(* IEC 61131-3 sources: STAR-PLC-Agent/results/raw/codex_matrix_resume_20261114/codex_deepseek/PUB019/functional/attempt_0001, 1 file *)

(* ---- test_program.st ---- *)
PROGRAM PLC_PRG
VAR
 BenchStep : UDINT := 0;
 BenchCalls : UDINT := 0;
 BenchDone : BOOL := FALSE;
 BenchUut0 : FB_Task;
 BenchUut1 : FB_Task;
 BenchUut2 : FB_Task;
 BenchUut3 : FB_Task;
 BenchUut4 : FB_Task;
 BenchUut5 : FB_Task;
 BenchUut6 : FB_Task;
 BenchUut7 : FB_Task;
 BenchUut8 : FB_Task;
 BenchUut9 : FB_Task;
 BenchUut10 : FB_Task;
 BenchUut11 : FB_Task;
 BenchUut12 : FB_Task;
 BenchUut13 : FB_Task;
 BenchUut14 : FB_Task;
 BenchUut15 : FB_Task;
 BenchUut16 : FB_Task;
 TraceIn_ManualMode : ARRAY[0..305] OF BOOL;
 TraceIn_SingleStepMode : ARRAY[0..305] OF BOOL;
 TraceIn_SingleCycleMode : ARRAY[0..305] OF BOOL;
 TraceIn_ContinuousMode : ARRAY[0..305] OF BOOL;
 TraceIn_EmergencyStop : ARRAY[0..305] OF BOOL;
 TraceIn_Start : ARRAY[0..305] OF BOOL;
 TraceIn_DownButton : ARRAY[0..305] OF BOOL;
 TraceIn_UpButton : ARRAY[0..305] OF BOOL;
 TraceIn_LeftButton : ARRAY[0..305] OF BOOL;
 TraceIn_RightButton : ARRAY[0..305] OF BOOL;
 TraceIn_GripButton : ARRAY[0..305] OF BOOL;
 TraceIn_ReleaseButton : ARRAY[0..305] OF BOOL;
 TraceIn_DownLimitSwitch : ARRAY[0..305] OF BOOL;
 TraceIn_UpLimitSwitch : ARRAY[0..305] OF BOOL;
 TraceIn_LeftLimitSwitch : ARRAY[0..305] OF BOOL;
 TraceIn_RightLimitSwitch : ARRAY[0..305] OF BOOL;
 TraceIn_GripLimitSwitch : ARRAY[0..305] OF BOOL;
 TraceIn_ReleaseLimitSwitch : ARRAY[0..305] OF BOOL;
 TraceOut_MoveDown : ARRAY[0..305] OF BOOL;
 TraceOut_MoveUp : ARRAY[0..305] OF BOOL;
 TraceOut_MoveLeft : ARRAY[0..305] OF BOOL;
 TraceOut_MoveRight : ARRAY[0..305] OF BOOL;
 TraceOut_ActivateGrip : ARRAY[0..305] OF BOOL;
 TraceOut_ActivateRelease : ARRAY[0..305] OF BOOL;
END_VAR

IF NOT BenchDone THEN
 CASE BenchStep OF
 0:
   BenchUut0.ManualMode := TRUE;
   BenchUut0.SingleStepMode := FALSE;
   BenchUut0.SingleCycleMode := FALSE;
   BenchUut0.ContinuousMode := FALSE;
   BenchUut0.EmergencyStop := TRUE;
   BenchUut0.Start := FALSE;
   BenchUut0.DownButton := TRUE;
   BenchUut0.UpButton := FALSE;
   BenchUut0.LeftButton := FALSE;
   BenchUut0.RightButton := FALSE;
   BenchUut0.GripButton := FALSE;
   BenchUut0.ReleaseButton := FALSE;
   BenchUut0.DownLimitSwitch := FALSE;
   BenchUut0.UpLimitSwitch := TRUE;
   BenchUut0.LeftLimitSwitch := TRUE;
   BenchUut0.RightLimitSwitch := FALSE;
   BenchUut0.GripLimitSwitch := FALSE;
   BenchUut0.ReleaseLimitSwitch := TRUE;
   TraceIn_ManualMode[0] := BenchUut0.ManualMode;
   TraceIn_SingleStepMode[0] := BenchUut0.SingleStepMode;
   TraceIn_SingleCycleMode[0] := BenchUut0.SingleCycleMode;
   TraceIn_ContinuousMode[0] := BenchUut0.ContinuousMode;
   TraceIn_EmergencyStop[0] := BenchUut0.EmergencyStop;
   TraceIn_Start[0] := BenchUut0.Start;
   TraceIn_DownButton[0] := BenchUut0.DownButton;
   TraceIn_UpButton[0] := BenchUut0.UpButton;
   TraceIn_LeftButton[0] := BenchUut0.LeftButton;
   TraceIn_RightButton[0] := BenchUut0.RightButton;
   TraceIn_GripButton[0] := BenchUut0.GripButton;
   TraceIn_ReleaseButton[0] := BenchUut0.ReleaseButton;
   TraceIn_DownLimitSwitch[0] := BenchUut0.DownLimitSwitch;
   TraceIn_UpLimitSwitch[0] := BenchUut0.UpLimitSwitch;
   TraceIn_LeftLimitSwitch[0] := BenchUut0.LeftLimitSwitch;
   TraceIn_RightLimitSwitch[0] := BenchUut0.RightLimitSwitch;
   TraceIn_GripLimitSwitch[0] := BenchUut0.GripLimitSwitch;
   TraceIn_ReleaseLimitSwitch[0] := BenchUut0.ReleaseLimitSwitch;
   BenchUut0();
   TraceOut_MoveDown[0] := BenchUut0.MoveDown;
   TraceOut_MoveUp[0] := BenchUut0.MoveUp;
   TraceOut_MoveLeft[0] := BenchUut0.MoveLeft;
   TraceOut_MoveRight[0] := BenchUut0.MoveRight;
   TraceOut_ActivateGrip[0] := BenchUut0.ActivateGrip;
   TraceOut_ActivateRelease[0] := BenchUut0.ActivateRelease;
   BenchCalls := BenchCalls + 1;
 1:
   BenchUut0.ManualMode := TRUE;
   BenchUut0.SingleStepMode := FALSE;
   BenchUut0.SingleCycleMode := FALSE;
   BenchUut0.ContinuousMode := FALSE;
   BenchUut0.EmergencyStop := TRUE;
   BenchUut0.Start := FALSE;
   BenchUut0.DownButton := TRUE;
   BenchUut0.UpButton := FALSE;
   BenchUut0.LeftButton := FALSE;
   BenchUut0.RightButton := FALSE;
   BenchUut0.GripButton := FALSE;
   BenchUut0.ReleaseButton := FALSE;
   BenchUut0.DownLimitSwitch := TRUE;
   BenchUut0.UpLimitSwitch := FALSE;
   BenchUut0.LeftLimitSwitch := TRUE;
   BenchUut0.RightLimitSwitch := FALSE;
   BenchUut0.GripLimitSwitch := FALSE;
   BenchUut0.ReleaseLimitSwitch := TRUE;
   TraceIn_ManualMode[1] := BenchUut0.ManualMode;
   TraceIn_SingleStepMode[1] := BenchUut0.SingleStepMode;
   TraceIn_SingleCycleMode[1] := BenchUut0.SingleCycleMode;
   TraceIn_ContinuousMode[1] := BenchUut0.ContinuousMode;
   TraceIn_EmergencyStop[1] := BenchUut0.EmergencyStop;
   TraceIn_Start[1] := BenchUut0.Start;
   TraceIn_DownButton[1] := BenchUut0.DownButton;
   TraceIn_UpButton[1] := BenchUut0.UpButton;
   TraceIn_LeftButton[1] := BenchUut0.LeftButton;
   TraceIn_RightButton[1] := BenchUut0.RightButton;
   TraceIn_GripButton[1] := BenchUut0.GripButton;
   TraceIn_ReleaseButton[1] := BenchUut0.ReleaseButton;
   TraceIn_DownLimitSwitch[1] := BenchUut0.DownLimitSwitch;
   TraceIn_UpLimitSwitch[1] := BenchUut0.UpLimitSwitch;
   TraceIn_LeftLimitSwitch[1] := BenchUut0.LeftLimitSwitch;
   TraceIn_RightLimitSwitch[1] := BenchUut0.RightLimitSwitch;
   TraceIn_GripLimitSwitch[1] := BenchUut0.GripLimitSwitch;
   TraceIn_ReleaseLimitSwitch[1] := BenchUut0.ReleaseLimitSwitch;
   BenchUut0();
   TraceOut_MoveDown[1] := BenchUut0.MoveDown;
   TraceOut_MoveUp[1] := BenchUut0.MoveUp;
   TraceOut_MoveLeft[1] := BenchUut0.MoveLeft;
   TraceOut_MoveRight[1] := BenchUut0.MoveRight;
   TraceOut_ActivateGrip[1] := BenchUut0.ActivateGrip;
   TraceOut_ActivateRelease[1] := BenchUut0.ActivateRelease;
   BenchCalls := BenchCalls + 1;
 2:
   BenchUut0.ManualMode := TRUE;
   BenchUut0.SingleStepMode := FALSE;
   BenchUut0.SingleCycleMode := FALSE;
   BenchUut0.ContinuousMode := FALSE;
   BenchUut0.EmergencyStop := TRUE;
   BenchUut0.Start := FALSE;
   BenchUut0.DownButton := FALSE;
   BenchUut0.UpButton := FALSE;
   BenchUut0.LeftButton := FALSE;
   BenchUut0.RightButton := FALSE;
   BenchUut0.GripButton := FALSE;
   BenchUut0.ReleaseButton := FALSE;
   BenchUut0.DownLimitSwitch := FALSE;
   BenchUut0.UpLimitSwitch := TRUE;
   BenchUut0.LeftLimitSwitch := TRUE;
   BenchUut0.RightLimitSwitch := FALSE;
   BenchUut0.GripLimitSwitch := FALSE;
   BenchUut0.ReleaseLimitSwitch := TRUE;
   TraceIn_ManualMode[2] := BenchUut0.ManualMode;
   TraceIn_SingleStepMode[2] := BenchUut0.SingleStepMode;
   TraceIn_SingleCycleMode[2] := BenchUut0.SingleCycleMode;
   TraceIn_ContinuousMode[2] := BenchUut0.ContinuousMode;
   TraceIn_EmergencyStop[2] := BenchUut0.EmergencyStop;
   TraceIn_Start[2] := BenchUut0.Start;
   TraceIn_DownButton[2] := BenchUut0.DownButton;
   TraceIn_UpButton[2] := BenchUut0.UpButton;
   TraceIn_LeftButton[2] := BenchUut0.LeftButton;
   TraceIn_RightButton[2] := BenchUut0.RightButton;
   TraceIn_GripButton[2] := BenchUut0.GripButton;
   TraceIn_ReleaseButton[2] := BenchUut0.ReleaseButton;
   TraceIn_DownLimitSwitch[2] := BenchUut0.DownLimitSwitch;
   TraceIn_UpLimitSwitch[2] := BenchUut0.UpLimitSwitch;
   TraceIn_LeftLimitSwitch[2] := BenchUut0.LeftLimitSwitch;
   TraceIn_RightLimitSwitch[2] := BenchUut0.RightLimitSwitch;
   TraceIn_GripLimitSwitch[2] := BenchUut0.GripLimitSwitch;
   TraceIn_ReleaseLimitSwitch[2] := BenchUut0.ReleaseLimitSwitch;
   BenchUut0();
   TraceOut_MoveDown[2] := BenchUut0.MoveDown;
   TraceOut_MoveUp[2] := BenchUut0.MoveUp;
   TraceOut_MoveLeft[2] := BenchUut0.MoveLeft;
   TraceOut_MoveRight[2] := BenchUut0.MoveRight;
   TraceOut_ActivateGrip[2] := BenchUut0.ActivateGrip;
   TraceOut_ActivateRelease[2] := BenchUut0.ActivateRelease;
   BenchCalls := BenchCalls + 1;
 3:
   BenchUut0.ManualMode := TRUE;
   BenchUut0.SingleStepMode := FALSE;
   BenchUut0.SingleCycleMode := FALSE;
   BenchUut0.ContinuousMode := FALSE;
   BenchUut0.EmergencyStop := TRUE;
   BenchUut0.Start := FALSE;
   BenchUut0.DownButton := TRUE;
   BenchUut0.UpButton := TRUE;
   BenchUut0.LeftButton := FALSE;
   BenchUut0.RightButton := FALSE;
   BenchUut0.GripButton := FALSE;
   BenchUut0.ReleaseButton := FALSE;
   BenchUut0.DownLimitSwitch := FALSE;
   BenchUut0.UpLimitSwitch := FALSE;
   BenchUut0.LeftLimitSwitch := TRUE;
   BenchUut0.RightLimitSwitch := FALSE;
   BenchUut0.GripLimitSwitch := FALSE;
   BenchUut0.ReleaseLimitSwitch := TRUE;
   TraceIn_ManualMode[3] := BenchUut0.ManualMode;
   TraceIn_SingleStepMode[3] := BenchUut0.SingleStepMode;
   TraceIn_SingleCycleMode[3] := BenchUut0.SingleCycleMode;
   TraceIn_ContinuousMode[3] := BenchUut0.ContinuousMode;
   TraceIn_EmergencyStop[3] := BenchUut0.EmergencyStop;
   TraceIn_Start[3] := BenchUut0.Start;
   TraceIn_DownButton[3] := BenchUut0.DownButton;
   TraceIn_UpButton[3] := BenchUut0.UpButton;
   TraceIn_LeftButton[3] := BenchUut0.LeftButton;
   TraceIn_RightButton[3] := BenchUut0.RightButton;
   TraceIn_GripButton[3] := BenchUut0.GripButton;
   TraceIn_ReleaseButton[3] := BenchUut0.ReleaseButton;
   TraceIn_DownLimitSwitch[3] := BenchUut0.DownLimitSwitch;
   TraceIn_UpLimitSwitch[3] := BenchUut0.UpLimitSwitch;
   TraceIn_LeftLimitSwitch[3] := BenchUut0.LeftLimitSwitch;
   TraceIn_RightLimitSwitch[3] := BenchUut0.RightLimitSwitch;
   TraceIn_GripLimitSwitch[3] := BenchUut0.GripLimitSwitch;
   TraceIn_ReleaseLimitSwitch[3] := BenchUut0.ReleaseLimitSwitch;
   BenchUut0();
   TraceOut_MoveDown[3] := BenchUut0.MoveDown;
   TraceOut_MoveUp[3] := BenchUut0.MoveUp;
   TraceOut_MoveLeft[3] := BenchUut0.MoveLeft;
   TraceOut_MoveRight[3] := BenchUut0.MoveRight;
   TraceOut_ActivateGrip[3] := BenchUut0.ActivateGrip;
   TraceOut_ActivateRelease[3] := BenchUut0.ActivateRelease;
   BenchCalls := BenchCalls + 1;
 4:
   BenchUut0.ManualMode := TRUE;
   BenchUut0.SingleStepMode := FALSE;
   BenchUut0.SingleCycleMode := FALSE;
   BenchUut0.ContinuousMode := FALSE;
   BenchUut0.EmergencyStop := TRUE;
   BenchUut0.Start := FALSE;
   BenchUut0.DownButton := FALSE;
   BenchUut0.UpButton := FALSE;
   BenchUut0.LeftButton := FALSE;
   BenchUut0.RightButton := TRUE;
   BenchUut0.GripButton := FALSE;
   BenchUut0.ReleaseButton := FALSE;
   BenchUut0.DownLimitSwitch := FALSE;
   BenchUut0.UpLimitSwitch := TRUE;
   BenchUut0.LeftLimitSwitch := TRUE;
   BenchUut0.RightLimitSwitch := FALSE;
   BenchUut0.GripLimitSwitch := FALSE;
   BenchUut0.ReleaseLimitSwitch := TRUE;
   TraceIn_ManualMode[4] := BenchUut0.ManualMode;
   TraceIn_SingleStepMode[4] := BenchUut0.SingleStepMode;
   TraceIn_SingleCycleMode[4] := BenchUut0.SingleCycleMode;
   TraceIn_ContinuousMode[4] := BenchUut0.ContinuousMode;
   TraceIn_EmergencyStop[4] := BenchUut0.EmergencyStop;
   TraceIn_Start[4] := BenchUut0.Start;
   TraceIn_DownButton[4] := BenchUut0.DownButton;
   TraceIn_UpButton[4] := BenchUut0.UpButton;
   TraceIn_LeftButton[4] := BenchUut0.LeftButton;
   TraceIn_RightButton[4] := BenchUut0.RightButton;
   TraceIn_GripButton[4] := BenchUut0.GripButton;
   TraceIn_ReleaseButton[4] := BenchUut0.ReleaseButton;
   TraceIn_DownLimitSwitch[4] := BenchUut0.DownLimitSwitch;
   TraceIn_UpLimitSwitch[4] := BenchUut0.UpLimitSwitch;
   TraceIn_LeftLimitSwitch[4] := BenchUut0.LeftLimitSwitch;
   TraceIn_RightLimitSwitch[4] := BenchUut0.RightLimitSwitch;
   TraceIn_GripLimitSwitch[4] := BenchUut0.GripLimitSwitch;
   TraceIn_ReleaseLimitSwitch[4] := BenchUut0.ReleaseLimitSwitch;
   BenchUut0();
   TraceOut_MoveDown[4] := BenchUut0.MoveDown;
   TraceOut_MoveUp[4] := BenchUut0.MoveUp;
   TraceOut_MoveLeft[4] := BenchUut0.MoveLeft;
   TraceOut_MoveRight[4] := BenchUut0.MoveRight;
   TraceOut_ActivateGrip[4] := BenchUut0.ActivateGrip;
   TraceOut_ActivateRelease[4] := BenchUut0.ActivateRelease;
   BenchCalls := BenchCalls + 1;
 5:
   BenchUut0.ManualMode := TRUE;
   BenchUut0.SingleStepMode := FALSE;
   BenchUut0.SingleCycleMode := FALSE;
   BenchUut0.ContinuousMode := FALSE;
   BenchUut0.EmergencyStop := TRUE;
   BenchUut0.Start := FALSE;
   BenchUut0.DownButton := FALSE;
   BenchUut0.UpButton := FALSE;
   BenchUut0.LeftButton := FALSE;
   BenchUut0.RightButton := TRUE;
   BenchUut0.GripButton := FALSE;
   BenchUut0.ReleaseButton := FALSE;
   BenchUut0.DownLimitSwitch := FALSE;
   BenchUut0.UpLimitSwitch := TRUE;
   BenchUut0.LeftLimitSwitch := FALSE;
   BenchUut0.RightLimitSwitch := TRUE;
   BenchUut0.GripLimitSwitch := FALSE;
   BenchUut0.ReleaseLimitSwitch := TRUE;
   TraceIn_ManualMode[5] := BenchUut0.ManualMode;
   TraceIn_SingleStepMode[5] := BenchUut0.SingleStepMode;
   TraceIn_SingleCycleMode[5] := BenchUut0.SingleCycleMode;
   TraceIn_ContinuousMode[5] := BenchUut0.ContinuousMode;
   TraceIn_EmergencyStop[5] := BenchUut0.EmergencyStop;
   TraceIn_Start[5] := BenchUut0.Start;
   TraceIn_DownButton[5] := BenchUut0.DownButton;
   TraceIn_UpButton[5] := BenchUut0.UpButton;
   TraceIn_LeftButton[5] := BenchUut0.LeftButton;
   TraceIn_RightButton[5] := BenchUut0.RightButton;
   TraceIn_GripButton[5] := BenchUut0.GripButton;
   TraceIn_ReleaseButton[5] := BenchUut0.ReleaseButton;
   TraceIn_DownLimitSwitch[5] := BenchUut0.DownLimitSwitch;
   TraceIn_UpLimitSwitch[5] := BenchUut0.UpLimitSwitch;
   TraceIn_LeftLimitSwitch[5] := BenchUut0.LeftLimitSwitch;
   TraceIn_RightLimitSwitch[5] := BenchUut0.RightLimitSwitch;
   TraceIn_GripLimitSwitch[5] := BenchUut0.GripLimitSwitch;
   TraceIn_ReleaseLimitSwitch[5] := BenchUut0.ReleaseLimitSwitch;
   BenchUut0();
   TraceOut_MoveDown[5] := BenchUut0.MoveDown;
   TraceOut_MoveUp[5] := BenchUut0.MoveUp;
   TraceOut_MoveLeft[5] := BenchUut0.MoveLeft;
   TraceOut_MoveRight[5] := BenchUut0.MoveRight;
   TraceOut_ActivateGrip[5] := BenchUut0.ActivateGrip;
   TraceOut_ActivateRelease[5] := BenchUut0.ActivateRelease;
   BenchCalls := BenchCalls + 1;
 6:
   BenchUut0.ManualMode := TRUE;
   BenchUut0.SingleStepMode := FALSE;
   BenchUut0.SingleCycleMode := FALSE;
   BenchUut0.ContinuousMode := FALSE;
   BenchUut0.EmergencyStop := TRUE;
   BenchUut0.Start := FALSE;
   BenchUut0.DownButton := FALSE;
   BenchUut0.UpButton := FALSE;
   BenchUut0.LeftButton := FALSE;
   BenchUut0.RightButton := FALSE;
   BenchUut0.GripButton := TRUE;
   BenchUut0.ReleaseButton := FALSE;
   BenchUut0.DownLimitSwitch := FALSE;
   BenchUut0.UpLimitSwitch := TRUE;
   BenchUut0.LeftLimitSwitch := TRUE;
   BenchUut0.RightLimitSwitch := FALSE;
   BenchUut0.GripLimitSwitch := FALSE;
   BenchUut0.ReleaseLimitSwitch := FALSE;
   TraceIn_ManualMode[6] := BenchUut0.ManualMode;
   TraceIn_SingleStepMode[6] := BenchUut0.SingleStepMode;
   TraceIn_SingleCycleMode[6] := BenchUut0.SingleCycleMode;
   TraceIn_ContinuousMode[6] := BenchUut0.ContinuousMode;
   TraceIn_EmergencyStop[6] := BenchUut0.EmergencyStop;
   TraceIn_Start[6] := BenchUut0.Start;
   TraceIn_DownButton[6] := BenchUut0.DownButton;
   TraceIn_UpButton[6] := BenchUut0.UpButton;
   TraceIn_LeftButton[6] := BenchUut0.LeftButton;
   TraceIn_RightButton[6] := BenchUut0.RightButton;
   TraceIn_GripButton[6] := BenchUut0.GripButton;
   TraceIn_ReleaseButton[6] := BenchUut0.ReleaseButton;
   TraceIn_DownLimitSwitch[6] := BenchUut0.DownLimitSwitch;
   TraceIn_UpLimitSwitch[6] := BenchUut0.UpLimitSwitch;
   TraceIn_LeftLimitSwitch[6] := BenchUut0.LeftLimitSwitch;
   TraceIn_RightLimitSwitch[6] := BenchUut0.RightLimitSwitch;
   TraceIn_GripLimitSwitch[6] := BenchUut0.GripLimitSwitch;
   TraceIn_ReleaseLimitSwitch[6] := BenchUut0.ReleaseLimitSwitch;
   BenchUut0();
   TraceOut_MoveDown[6] := BenchUut0.MoveDown;
   TraceOut_MoveUp[6] := BenchUut0.MoveUp;
   TraceOut_MoveLeft[6] := BenchUut0.MoveLeft;
   TraceOut_MoveRight[6] := BenchUut0.MoveRight;
   TraceOut_ActivateGrip[6] := BenchUut0.ActivateGrip;
   TraceOut_ActivateRelease[6] := BenchUut0.ActivateRelease;
   BenchCalls := BenchCalls + 1;
 7:
   BenchUut0.ManualMode := TRUE;
   BenchUut0.SingleStepMode := FALSE;
   BenchUut0.SingleCycleMode := FALSE;
   BenchUut0.ContinuousMode := FALSE;
   BenchUut0.EmergencyStop := TRUE;
   BenchUut0.Start := FALSE;
   BenchUut0.DownButton := FALSE;
   BenchUut0.UpButton := FALSE;
   BenchUut0.LeftButton := FALSE;
   BenchUut0.RightButton := FALSE;
   BenchUut0.GripButton := TRUE;
   BenchUut0.ReleaseButton := FALSE;
   BenchUut0.DownLimitSwitch := FALSE;
   BenchUut0.UpLimitSwitch := TRUE;
   BenchUut0.LeftLimitSwitch := TRUE;
   BenchUut0.RightLimitSwitch := FALSE;
   BenchUut0.GripLimitSwitch := TRUE;
   BenchUut0.ReleaseLimitSwitch := FALSE;
   TraceIn_ManualMode[7] := BenchUut0.ManualMode;
   TraceIn_SingleStepMode[7] := BenchUut0.SingleStepMode;
   TraceIn_SingleCycleMode[7] := BenchUut0.SingleCycleMode;
   TraceIn_ContinuousMode[7] := BenchUut0.ContinuousMode;
   TraceIn_EmergencyStop[7] := BenchUut0.EmergencyStop;
   TraceIn_Start[7] := BenchUut0.Start;
   TraceIn_DownButton[7] := BenchUut0.DownButton;
   TraceIn_UpButton[7] := BenchUut0.UpButton;
   TraceIn_LeftButton[7] := BenchUut0.LeftButton;
   TraceIn_RightButton[7] := BenchUut0.RightButton;
   TraceIn_GripButton[7] := BenchUut0.GripButton;
   TraceIn_ReleaseButton[7] := BenchUut0.ReleaseButton;
   TraceIn_DownLimitSwitch[7] := BenchUut0.DownLimitSwitch;
   TraceIn_UpLimitSwitch[7] := BenchUut0.UpLimitSwitch;
   TraceIn_LeftLimitSwitch[7] := BenchUut0.LeftLimitSwitch;
   TraceIn_RightLimitSwitch[7] := BenchUut0.RightLimitSwitch;
   TraceIn_GripLimitSwitch[7] := BenchUut0.GripLimitSwitch;
   TraceIn_ReleaseLimitSwitch[7] := BenchUut0.ReleaseLimitSwitch;
   BenchUut0();
   TraceOut_MoveDown[7] := BenchUut0.MoveDown;
   TraceOut_MoveUp[7] := BenchUut0.MoveUp;
   TraceOut_MoveLeft[7] := BenchUut0.MoveLeft;
   TraceOut_MoveRight[7] := BenchUut0.MoveRight;
   TraceOut_ActivateGrip[7] := BenchUut0.ActivateGrip;
   TraceOut_ActivateRelease[7] := BenchUut0.ActivateRelease;
   BenchCalls := BenchCalls + 1;
 8:
   BenchUut0.ManualMode := TRUE;
   BenchUut0.SingleStepMode := FALSE;
   BenchUut0.SingleCycleMode := FALSE;
   BenchUut0.ContinuousMode := FALSE;
   BenchUut0.EmergencyStop := TRUE;
   BenchUut0.Start := FALSE;
   BenchUut0.DownButton := FALSE;
   BenchUut0.UpButton := FALSE;
   BenchUut0.LeftButton := FALSE;
   BenchUut0.RightButton := FALSE;
   BenchUut0.GripButton := TRUE;
   BenchUut0.ReleaseButton := TRUE;
   BenchUut0.DownLimitSwitch := FALSE;
   BenchUut0.UpLimitSwitch := TRUE;
   BenchUut0.LeftLimitSwitch := TRUE;
   BenchUut0.RightLimitSwitch := FALSE;
   BenchUut0.GripLimitSwitch := FALSE;
   BenchUut0.ReleaseLimitSwitch := FALSE;
   TraceIn_ManualMode[8] := BenchUut0.ManualMode;
   TraceIn_SingleStepMode[8] := BenchUut0.SingleStepMode;
   TraceIn_SingleCycleMode[8] := BenchUut0.SingleCycleMode;
   TraceIn_ContinuousMode[8] := BenchUut0.ContinuousMode;
   TraceIn_EmergencyStop[8] := BenchUut0.EmergencyStop;
   TraceIn_Start[8] := BenchUut0.Start;
   TraceIn_DownButton[8] := BenchUut0.DownButton;
   TraceIn_UpButton[8] := BenchUut0.UpButton;
   TraceIn_LeftButton[8] := BenchUut0.LeftButton;
   TraceIn_RightButton[8] := BenchUut0.RightButton;
   TraceIn_GripButton[8] := BenchUut0.GripButton;
   TraceIn_ReleaseButton[8] := BenchUut0.ReleaseButton;
   TraceIn_DownLimitSwitch[8] := BenchUut0.DownLimitSwitch;
   TraceIn_UpLimitSwitch[8] := BenchUut0.UpLimitSwitch;
   TraceIn_LeftLimitSwitch[8] := BenchUut0.LeftLimitSwitch;
   TraceIn_RightLimitSwitch[8] := BenchUut0.RightLimitSwitch;
   TraceIn_GripLimitSwitch[8] := BenchUut0.GripLimitSwitch;
   TraceIn_ReleaseLimitSwitch[8] := BenchUut0.ReleaseLimitSwitch;
   BenchUut0();
   TraceOut_MoveDown[8] := BenchUut0.MoveDown;
   TraceOut_MoveUp[8] := BenchUut0.MoveUp;
   TraceOut_MoveLeft[8] := BenchUut0.MoveLeft;
   TraceOut_MoveRight[8] := BenchUut0.MoveRight;
   TraceOut_ActivateGrip[8] := BenchUut0.ActivateGrip;
   TraceOut_ActivateRelease[8] := BenchUut0.ActivateRelease;
   BenchCalls := BenchCalls + 1;
 9:
   BenchUut0.ManualMode := TRUE;
   BenchUut0.SingleStepMode := FALSE;
   BenchUut0.SingleCycleMode := FALSE;
   BenchUut0.ContinuousMode := FALSE;
   BenchUut0.EmergencyStop := FALSE;
   BenchUut0.Start := FALSE;
   BenchUut0.DownButton := TRUE;
   BenchUut0.UpButton := FALSE;
   BenchUut0.LeftButton := FALSE;
   BenchUut0.RightButton := TRUE;
   BenchUut0.GripButton := FALSE;
   BenchUut0.ReleaseButton := FALSE;
   BenchUut0.DownLimitSwitch := FALSE;
   BenchUut0.UpLimitSwitch := TRUE;
   BenchUut0.LeftLimitSwitch := TRUE;
   BenchUut0.RightLimitSwitch := FALSE;
   BenchUut0.GripLimitSwitch := FALSE;
   BenchUut0.ReleaseLimitSwitch := TRUE;
   TraceIn_ManualMode[9] := BenchUut0.ManualMode;
   TraceIn_SingleStepMode[9] := BenchUut0.SingleStepMode;
   TraceIn_SingleCycleMode[9] := BenchUut0.SingleCycleMode;
   TraceIn_ContinuousMode[9] := BenchUut0.ContinuousMode;
   TraceIn_EmergencyStop[9] := BenchUut0.EmergencyStop;
   TraceIn_Start[9] := BenchUut0.Start;
   TraceIn_DownButton[9] := BenchUut0.DownButton;
   TraceIn_UpButton[9] := BenchUut0.UpButton;
   TraceIn_LeftButton[9] := BenchUut0.LeftButton;
   TraceIn_RightButton[9] := BenchUut0.RightButton;
   TraceIn_GripButton[9] := BenchUut0.GripButton;
   TraceIn_ReleaseButton[9] := BenchUut0.ReleaseButton;
   TraceIn_DownLimitSwitch[9] := BenchUut0.DownLimitSwitch;
   TraceIn_UpLimitSwitch[9] := BenchUut0.UpLimitSwitch;
   TraceIn_LeftLimitSwitch[9] := BenchUut0.LeftLimitSwitch;
   TraceIn_RightLimitSwitch[9] := BenchUut0.RightLimitSwitch;
   TraceIn_GripLimitSwitch[9] := BenchUut0.GripLimitSwitch;
   TraceIn_ReleaseLimitSwitch[9] := BenchUut0.ReleaseLimitSwitch;
   BenchUut0();
   TraceOut_MoveDown[9] := BenchUut0.MoveDown;
   TraceOut_MoveUp[9] := BenchUut0.MoveUp;
   TraceOut_MoveLeft[9] := BenchUut0.MoveLeft;
   TraceOut_MoveRight[9] := BenchUut0.MoveRight;
   TraceOut_ActivateGrip[9] := BenchUut0.ActivateGrip;
   TraceOut_ActivateRelease[9] := BenchUut0.ActivateRelease;
   BenchCalls := BenchCalls + 1;
 10:
   BenchUut1.ManualMode := FALSE;
   BenchUut1.SingleStepMode := TRUE;
   BenchUut1.SingleCycleMode := FALSE;
   BenchUut1.ContinuousMode := FALSE;
   BenchUut1.EmergencyStop := TRUE;
   BenchUut1.Start := FALSE;
   BenchUut1.DownButton := FALSE;
   BenchUut1.UpButton := FALSE;
   BenchUut1.LeftButton := FALSE;
   BenchUut1.RightButton := FALSE;
   BenchUut1.GripButton := FALSE;
   BenchUut1.ReleaseButton := FALSE;
   BenchUut1.DownLimitSwitch := FALSE;
   BenchUut1.UpLimitSwitch := TRUE;
   BenchUut1.LeftLimitSwitch := TRUE;
   BenchUut1.RightLimitSwitch := FALSE;
   BenchUut1.GripLimitSwitch := FALSE;
   BenchUut1.ReleaseLimitSwitch := TRUE;
   TraceIn_ManualMode[10] := BenchUut1.ManualMode;
   TraceIn_SingleStepMode[10] := BenchUut1.SingleStepMode;
   TraceIn_SingleCycleMode[10] := BenchUut1.SingleCycleMode;
   TraceIn_ContinuousMode[10] := BenchUut1.ContinuousMode;
   TraceIn_EmergencyStop[10] := BenchUut1.EmergencyStop;
   TraceIn_Start[10] := BenchUut1.Start;
   TraceIn_DownButton[10] := BenchUut1.DownButton;
   TraceIn_UpButton[10] := BenchUut1.UpButton;
   TraceIn_LeftButton[10] := BenchUut1.LeftButton;
   TraceIn_RightButton[10] := BenchUut1.RightButton;
   TraceIn_GripButton[10] := BenchUut1.GripButton;
   TraceIn_ReleaseButton[10] := BenchUut1.ReleaseButton;
   TraceIn_DownLimitSwitch[10] := BenchUut1.DownLimitSwitch;
   TraceIn_UpLimitSwitch[10] := BenchUut1.UpLimitSwitch;
   TraceIn_LeftLimitSwitch[10] := BenchUut1.LeftLimitSwitch;
   TraceIn_RightLimitSwitch[10] := BenchUut1.RightLimitSwitch;
   TraceIn_GripLimitSwitch[10] := BenchUut1.GripLimitSwitch;
   TraceIn_ReleaseLimitSwitch[10] := BenchUut1.ReleaseLimitSwitch;
   BenchUut1();
   TraceOut_MoveDown[10] := BenchUut1.MoveDown;
   TraceOut_MoveUp[10] := BenchUut1.MoveUp;
   TraceOut_MoveLeft[10] := BenchUut1.MoveLeft;
   TraceOut_MoveRight[10] := BenchUut1.MoveRight;
   TraceOut_ActivateGrip[10] := BenchUut1.ActivateGrip;
   TraceOut_ActivateRelease[10] := BenchUut1.ActivateRelease;
   BenchCalls := BenchCalls + 1;
 11:
   BenchUut1.ManualMode := FALSE;
   BenchUut1.SingleStepMode := TRUE;
   BenchUut1.SingleCycleMode := FALSE;
   BenchUut1.ContinuousMode := FALSE;
   BenchUut1.EmergencyStop := TRUE;
   BenchUut1.Start := TRUE;
   BenchUut1.DownButton := FALSE;
   BenchUut1.UpButton := FALSE;
   BenchUut1.LeftButton := FALSE;
   BenchUut1.RightButton := FALSE;
   BenchUut1.GripButton := FALSE;
   BenchUut1.ReleaseButton := FALSE;
   BenchUut1.DownLimitSwitch := FALSE;
   BenchUut1.UpLimitSwitch := TRUE;
   BenchUut1.LeftLimitSwitch := TRUE;
   BenchUut1.RightLimitSwitch := FALSE;
   BenchUut1.GripLimitSwitch := FALSE;
   BenchUut1.ReleaseLimitSwitch := TRUE;
   TraceIn_ManualMode[11] := BenchUut1.ManualMode;
   TraceIn_SingleStepMode[11] := BenchUut1.SingleStepMode;
   TraceIn_SingleCycleMode[11] := BenchUut1.SingleCycleMode;
   TraceIn_ContinuousMode[11] := BenchUut1.ContinuousMode;
   TraceIn_EmergencyStop[11] := BenchUut1.EmergencyStop;
   TraceIn_Start[11] := BenchUut1.Start;
   TraceIn_DownButton[11] := BenchUut1.DownButton;
   TraceIn_UpButton[11] := BenchUut1.UpButton;
   TraceIn_LeftButton[11] := BenchUut1.LeftButton;
   TraceIn_RightButton[11] := BenchUut1.RightButton;
   TraceIn_GripButton[11] := BenchUut1.GripButton;
   TraceIn_ReleaseButton[11] := BenchUut1.ReleaseButton;
   TraceIn_DownLimitSwitch[11] := BenchUut1.DownLimitSwitch;
   TraceIn_UpLimitSwitch[11] := BenchUut1.UpLimitSwitch;
   TraceIn_LeftLimitSwitch[11] := BenchUut1.LeftLimitSwitch;
   TraceIn_RightLimitSwitch[11] := BenchUut1.RightLimitSwitch;
   TraceIn_GripLimitSwitch[11] := BenchUut1.GripLimitSwitch;
   TraceIn_ReleaseLimitSwitch[11] := BenchUut1.ReleaseLimitSwitch;
   BenchUut1();
   TraceOut_MoveDown[11] := BenchUut1.MoveDown;
   TraceOut_MoveUp[11] := BenchUut1.MoveUp;
   TraceOut_MoveLeft[11] := BenchUut1.MoveLeft;
   TraceOut_MoveRight[11] := BenchUut1.MoveRight;
   TraceOut_ActivateGrip[11] := BenchUut1.ActivateGrip;
   TraceOut_ActivateRelease[11] := BenchUut1.ActivateRelease;
   BenchCalls := BenchCalls + 1;
 12:
   BenchUut1.ManualMode := FALSE;
   BenchUut1.SingleStepMode := TRUE;
   BenchUut1.SingleCycleMode := FALSE;
   BenchUut1.ContinuousMode := FALSE;
   BenchUut1.EmergencyStop := TRUE;
   BenchUut1.Start := TRUE;
   BenchUut1.DownButton := FALSE;
   BenchUut1.UpButton := FALSE;
   BenchUut1.LeftButton := FALSE;
   BenchUut1.RightButton := FALSE;
   BenchUut1.GripButton := FALSE;
   BenchUut1.ReleaseButton := FALSE;
   BenchUut1.DownLimitSwitch := FALSE;
   BenchUut1.UpLimitSwitch := FALSE;
   BenchUut1.LeftLimitSwitch := TRUE;
   BenchUut1.RightLimitSwitch := FALSE;
   BenchUut1.GripLimitSwitch := FALSE;
   BenchUut1.ReleaseLimitSwitch := TRUE;
   TraceIn_ManualMode[12] := BenchUut1.ManualMode;
   TraceIn_SingleStepMode[12] := BenchUut1.SingleStepMode;
   TraceIn_SingleCycleMode[12] := BenchUut1.SingleCycleMode;
   TraceIn_ContinuousMode[12] := BenchUut1.ContinuousMode;
   TraceIn_EmergencyStop[12] := BenchUut1.EmergencyStop;
   TraceIn_Start[12] := BenchUut1.Start;
   TraceIn_DownButton[12] := BenchUut1.DownButton;
   TraceIn_UpButton[12] := BenchUut1.UpButton;
   TraceIn_LeftButton[12] := BenchUut1.LeftButton;
   TraceIn_RightButton[12] := BenchUut1.RightButton;
   TraceIn_GripButton[12] := BenchUut1.GripButton;
   TraceIn_ReleaseButton[12] := BenchUut1.ReleaseButton;
   TraceIn_DownLimitSwitch[12] := BenchUut1.DownLimitSwitch;
   TraceIn_UpLimitSwitch[12] := BenchUut1.UpLimitSwitch;
   TraceIn_LeftLimitSwitch[12] := BenchUut1.LeftLimitSwitch;
   TraceIn_RightLimitSwitch[12] := BenchUut1.RightLimitSwitch;
   TraceIn_GripLimitSwitch[12] := BenchUut1.GripLimitSwitch;
   TraceIn_ReleaseLimitSwitch[12] := BenchUut1.ReleaseLimitSwitch;
   BenchUut1();
   TraceOut_MoveDown[12] := BenchUut1.MoveDown;
   TraceOut_MoveUp[12] := BenchUut1.MoveUp;
   TraceOut_MoveLeft[12] := BenchUut1.MoveLeft;
   TraceOut_MoveRight[12] := BenchUut1.MoveRight;
   TraceOut_ActivateGrip[12] := BenchUut1.ActivateGrip;
   TraceOut_ActivateRelease[12] := BenchUut1.ActivateRelease;
   BenchCalls := BenchCalls + 1;
 13:
   BenchUut1.ManualMode := FALSE;
   BenchUut1.SingleStepMode := TRUE;
   BenchUut1.SingleCycleMode := FALSE;
   BenchUut1.ContinuousMode := FALSE;
   BenchUut1.EmergencyStop := TRUE;
   BenchUut1.Start := TRUE;
   BenchUut1.DownButton := FALSE;
   BenchUut1.UpButton := FALSE;
   BenchUut1.LeftButton := FALSE;
   BenchUut1.RightButton := FALSE;
   BenchUut1.GripButton := FALSE;
   BenchUut1.ReleaseButton := FALSE;
   BenchUut1.DownLimitSwitch := TRUE;
   BenchUut1.UpLimitSwitch := FALSE;
   BenchUut1.LeftLimitSwitch := TRUE;
   BenchUut1.RightLimitSwitch := FALSE;
   BenchUut1.GripLimitSwitch := FALSE;
   BenchUut1.ReleaseLimitSwitch := TRUE;
   TraceIn_ManualMode[13] := BenchUut1.ManualMode;
   TraceIn_SingleStepMode[13] := BenchUut1.SingleStepMode;
   TraceIn_SingleCycleMode[13] := BenchUut1.SingleCycleMode;
   TraceIn_ContinuousMode[13] := BenchUut1.ContinuousMode;
   TraceIn_EmergencyStop[13] := BenchUut1.EmergencyStop;
   TraceIn_Start[13] := BenchUut1.Start;
   TraceIn_DownButton[13] := BenchUut1.DownButton;
   TraceIn_UpButton[13] := BenchUut1.UpButton;
   TraceIn_LeftButton[13] := BenchUut1.LeftButton;
   TraceIn_RightButton[13] := BenchUut1.RightButton;
   TraceIn_GripButton[13] := BenchUut1.GripButton;
   TraceIn_ReleaseButton[13] := BenchUut1.ReleaseButton;
   TraceIn_DownLimitSwitch[13] := BenchUut1.DownLimitSwitch;
   TraceIn_UpLimitSwitch[13] := BenchUut1.UpLimitSwitch;
   TraceIn_LeftLimitSwitch[13] := BenchUut1.LeftLimitSwitch;
   TraceIn_RightLimitSwitch[13] := BenchUut1.RightLimitSwitch;
   TraceIn_GripLimitSwitch[13] := BenchUut1.GripLimitSwitch;
   TraceIn_ReleaseLimitSwitch[13] := BenchUut1.ReleaseLimitSwitch;
   BenchUut1();
   TraceOut_MoveDown[13] := BenchUut1.MoveDown;
   TraceOut_MoveUp[13] := BenchUut1.MoveUp;
   TraceOut_MoveLeft[13] := BenchUut1.MoveLeft;
   TraceOut_MoveRight[13] := BenchUut1.MoveRight;
   TraceOut_ActivateGrip[13] := BenchUut1.ActivateGrip;
   TraceOut_ActivateRelease[13] := BenchUut1.ActivateRelease;
   BenchCalls := BenchCalls + 1;
 14:
   BenchUut1.ManualMode := FALSE;
   BenchUut1.SingleStepMode := TRUE;
   BenchUut1.SingleCycleMode := FALSE;
   BenchUut1.ContinuousMode := FALSE;
   BenchUut1.EmergencyStop := TRUE;
   BenchUut1.Start := TRUE;
   BenchUut1.DownButton := FALSE;
   BenchUut1.UpButton := FALSE;
   BenchUut1.LeftButton := FALSE;
   BenchUut1.RightButton := FALSE;
   BenchUut1.GripButton := FALSE;
   BenchUut1.ReleaseButton := FALSE;
   BenchUut1.DownLimitSwitch := TRUE;
   BenchUut1.UpLimitSwitch := FALSE;
   BenchUut1.LeftLimitSwitch := TRUE;
   BenchUut1.RightLimitSwitch := FALSE;
   BenchUut1.GripLimitSwitch := FALSE;
   BenchUut1.ReleaseLimitSwitch := TRUE;
   TraceIn_ManualMode[14] := BenchUut1.ManualMode;
   TraceIn_SingleStepMode[14] := BenchUut1.SingleStepMode;
   TraceIn_SingleCycleMode[14] := BenchUut1.SingleCycleMode;
   TraceIn_ContinuousMode[14] := BenchUut1.ContinuousMode;
   TraceIn_EmergencyStop[14] := BenchUut1.EmergencyStop;
   TraceIn_Start[14] := BenchUut1.Start;
   TraceIn_DownButton[14] := BenchUut1.DownButton;
   TraceIn_UpButton[14] := BenchUut1.UpButton;
   TraceIn_LeftButton[14] := BenchUut1.LeftButton;
   TraceIn_RightButton[14] := BenchUut1.RightButton;
   TraceIn_GripButton[14] := BenchUut1.GripButton;
   TraceIn_ReleaseButton[14] := BenchUut1.ReleaseButton;
   TraceIn_DownLimitSwitch[14] := BenchUut1.DownLimitSwitch;
   TraceIn_UpLimitSwitch[14] := BenchUut1.UpLimitSwitch;
   TraceIn_LeftLimitSwitch[14] := BenchUut1.LeftLimitSwitch;
   TraceIn_RightLimitSwitch[14] := BenchUut1.RightLimitSwitch;
   TraceIn_GripLimitSwitch[14] := BenchUut1.GripLimitSwitch;
   TraceIn_ReleaseLimitSwitch[14] := BenchUut1.ReleaseLimitSwitch;
   BenchUut1();
   TraceOut_MoveDown[14] := BenchUut1.MoveDown;
   TraceOut_MoveUp[14] := BenchUut1.MoveUp;
   TraceOut_MoveLeft[14] := BenchUut1.MoveLeft;
   TraceOut_MoveRight[14] := BenchUut1.MoveRight;
   TraceOut_ActivateGrip[14] := BenchUut1.ActivateGrip;
   TraceOut_ActivateRelease[14] := BenchUut1.ActivateRelease;
   BenchCalls := BenchCalls + 1;
 15:
   BenchUut1.ManualMode := FALSE;
   BenchUut1.SingleStepMode := TRUE;
   BenchUut1.SingleCycleMode := FALSE;
   BenchUut1.ContinuousMode := FALSE;
   BenchUut1.EmergencyStop := TRUE;
   BenchUut1.Start := FALSE;
   BenchUut1.DownButton := FALSE;
   BenchUut1.UpButton := FALSE;
   BenchUut1.LeftButton := FALSE;
   BenchUut1.RightButton := FALSE;
   BenchUut1.GripButton := FALSE;
   BenchUut1.ReleaseButton := FALSE;
   BenchUut1.DownLimitSwitch := TRUE;
   BenchUut1.UpLimitSwitch := FALSE;
   BenchUut1.LeftLimitSwitch := TRUE;
   BenchUut1.RightLimitSwitch := FALSE;
   BenchUut1.GripLimitSwitch := FALSE;
   BenchUut1.ReleaseLimitSwitch := TRUE;
   TraceIn_ManualMode[15] := BenchUut1.ManualMode;
   TraceIn_SingleStepMode[15] := BenchUut1.SingleStepMode;
   TraceIn_SingleCycleMode[15] := BenchUut1.SingleCycleMode;
   TraceIn_ContinuousMode[15] := BenchUut1.ContinuousMode;
   TraceIn_EmergencyStop[15] := BenchUut1.EmergencyStop;
   TraceIn_Start[15] := BenchUut1.Start;
   TraceIn_DownButton[15] := BenchUut1.DownButton;
   TraceIn_UpButton[15] := BenchUut1.UpButton;
   TraceIn_LeftButton[15] := BenchUut1.LeftButton;
   TraceIn_RightButton[15] := BenchUut1.RightButton;
   TraceIn_GripButton[15] := BenchUut1.GripButton;
   TraceIn_ReleaseButton[15] := BenchUut1.ReleaseButton;
   TraceIn_DownLimitSwitch[15] := BenchUut1.DownLimitSwitch;
   TraceIn_UpLimitSwitch[15] := BenchUut1.UpLimitSwitch;
   TraceIn_LeftLimitSwitch[15] := BenchUut1.LeftLimitSwitch;
   TraceIn_RightLimitSwitch[15] := BenchUut1.RightLimitSwitch;
   TraceIn_GripLimitSwitch[15] := BenchUut1.GripLimitSwitch;
   TraceIn_ReleaseLimitSwitch[15] := BenchUut1.ReleaseLimitSwitch;
   BenchUut1();
   TraceOut_MoveDown[15] := BenchUut1.MoveDown;
   TraceOut_MoveUp[15] := BenchUut1.MoveUp;
   TraceOut_MoveLeft[15] := BenchUut1.MoveLeft;
   TraceOut_MoveRight[15] := BenchUut1.MoveRight;
   TraceOut_ActivateGrip[15] := BenchUut1.ActivateGrip;
   TraceOut_ActivateRelease[15] := BenchUut1.ActivateRelease;
   BenchCalls := BenchCalls + 1;
 16:
   BenchUut1.ManualMode := FALSE;
   BenchUut1.SingleStepMode := TRUE;
   BenchUut1.SingleCycleMode := FALSE;
   BenchUut1.ContinuousMode := FALSE;
   BenchUut1.EmergencyStop := TRUE;
   BenchUut1.Start := TRUE;
   BenchUut1.DownButton := FALSE;
   BenchUut1.UpButton := FALSE;
   BenchUut1.LeftButton := FALSE;
   BenchUut1.RightButton := FALSE;
   BenchUut1.GripButton := FALSE;
   BenchUut1.ReleaseButton := FALSE;
   BenchUut1.DownLimitSwitch := TRUE;
   BenchUut1.UpLimitSwitch := FALSE;
   BenchUut1.LeftLimitSwitch := TRUE;
   BenchUut1.RightLimitSwitch := FALSE;
   BenchUut1.GripLimitSwitch := FALSE;
   BenchUut1.ReleaseLimitSwitch := FALSE;
   TraceIn_ManualMode[16] := BenchUut1.ManualMode;
   TraceIn_SingleStepMode[16] := BenchUut1.SingleStepMode;
   TraceIn_SingleCycleMode[16] := BenchUut1.SingleCycleMode;
   TraceIn_ContinuousMode[16] := BenchUut1.ContinuousMode;
   TraceIn_EmergencyStop[16] := BenchUut1.EmergencyStop;
   TraceIn_Start[16] := BenchUut1.Start;
   TraceIn_DownButton[16] := BenchUut1.DownButton;
   TraceIn_UpButton[16] := BenchUut1.UpButton;
   TraceIn_LeftButton[16] := BenchUut1.LeftButton;
   TraceIn_RightButton[16] := BenchUut1.RightButton;
   TraceIn_GripButton[16] := BenchUut1.GripButton;
   TraceIn_ReleaseButton[16] := BenchUut1.ReleaseButton;
   TraceIn_DownLimitSwitch[16] := BenchUut1.DownLimitSwitch;
   TraceIn_UpLimitSwitch[16] := BenchUut1.UpLimitSwitch;
   TraceIn_LeftLimitSwitch[16] := BenchUut1.LeftLimitSwitch;
   TraceIn_RightLimitSwitch[16] := BenchUut1.RightLimitSwitch;
   TraceIn_GripLimitSwitch[16] := BenchUut1.GripLimitSwitch;
   TraceIn_ReleaseLimitSwitch[16] := BenchUut1.ReleaseLimitSwitch;
   BenchUut1();
   TraceOut_MoveDown[16] := BenchUut1.MoveDown;
   TraceOut_MoveUp[16] := BenchUut1.MoveUp;
   TraceOut_MoveLeft[16] := BenchUut1.MoveLeft;
   TraceOut_MoveRight[16] := BenchUut1.MoveRight;
   TraceOut_ActivateGrip[16] := BenchUut1.ActivateGrip;
   TraceOut_ActivateRelease[16] := BenchUut1.ActivateRelease;
   BenchCalls := BenchCalls + 1;
 17:
   BenchUut1.ManualMode := FALSE;
   BenchUut1.SingleStepMode := TRUE;
   BenchUut1.SingleCycleMode := FALSE;
   BenchUut1.ContinuousMode := FALSE;
   BenchUut1.EmergencyStop := TRUE;
   BenchUut1.Start := FALSE;
   BenchUut1.DownButton := FALSE;
   BenchUut1.UpButton := FALSE;
   BenchUut1.LeftButton := FALSE;
   BenchUut1.RightButton := FALSE;
   BenchUut1.GripButton := FALSE;
   BenchUut1.ReleaseButton := FALSE;
   BenchUut1.DownLimitSwitch := TRUE;
   BenchUut1.UpLimitSwitch := FALSE;
   BenchUut1.LeftLimitSwitch := TRUE;
   BenchUut1.RightLimitSwitch := FALSE;
   BenchUut1.GripLimitSwitch := TRUE;
   BenchUut1.ReleaseLimitSwitch := FALSE;
   TraceIn_ManualMode[17] := BenchUut1.ManualMode;
   TraceIn_SingleStepMode[17] := BenchUut1.SingleStepMode;
   TraceIn_SingleCycleMode[17] := BenchUut1.SingleCycleMode;
   TraceIn_ContinuousMode[17] := BenchUut1.ContinuousMode;
   TraceIn_EmergencyStop[17] := BenchUut1.EmergencyStop;
   TraceIn_Start[17] := BenchUut1.Start;
   TraceIn_DownButton[17] := BenchUut1.DownButton;
   TraceIn_UpButton[17] := BenchUut1.UpButton;
   TraceIn_LeftButton[17] := BenchUut1.LeftButton;
   TraceIn_RightButton[17] := BenchUut1.RightButton;
   TraceIn_GripButton[17] := BenchUut1.GripButton;
   TraceIn_ReleaseButton[17] := BenchUut1.ReleaseButton;
   TraceIn_DownLimitSwitch[17] := BenchUut1.DownLimitSwitch;
   TraceIn_UpLimitSwitch[17] := BenchUut1.UpLimitSwitch;
   TraceIn_LeftLimitSwitch[17] := BenchUut1.LeftLimitSwitch;
   TraceIn_RightLimitSwitch[17] := BenchUut1.RightLimitSwitch;
   TraceIn_GripLimitSwitch[17] := BenchUut1.GripLimitSwitch;
   TraceIn_ReleaseLimitSwitch[17] := BenchUut1.ReleaseLimitSwitch;
   BenchUut1();
   TraceOut_MoveDown[17] := BenchUut1.MoveDown;
   TraceOut_MoveUp[17] := BenchUut1.MoveUp;
   TraceOut_MoveLeft[17] := BenchUut1.MoveLeft;
   TraceOut_MoveRight[17] := BenchUut1.MoveRight;
   TraceOut_ActivateGrip[17] := BenchUut1.ActivateGrip;
   TraceOut_ActivateRelease[17] := BenchUut1.ActivateRelease;
   BenchCalls := BenchCalls + 1;
 18:
   BenchUut1.ManualMode := FALSE;
   BenchUut1.SingleStepMode := TRUE;
   BenchUut1.SingleCycleMode := FALSE;
   BenchUut1.ContinuousMode := FALSE;
   BenchUut1.EmergencyStop := TRUE;
   BenchUut1.Start := TRUE;
   BenchUut1.DownButton := FALSE;
   BenchUut1.UpButton := FALSE;
   BenchUut1.LeftButton := FALSE;
   BenchUut1.RightButton := FALSE;
   BenchUut1.GripButton := FALSE;
   BenchUut1.ReleaseButton := FALSE;
   BenchUut1.DownLimitSwitch := TRUE;
   BenchUut1.UpLimitSwitch := FALSE;
   BenchUut1.LeftLimitSwitch := TRUE;
   BenchUut1.RightLimitSwitch := FALSE;
   BenchUut1.GripLimitSwitch := TRUE;
   BenchUut1.ReleaseLimitSwitch := FALSE;
   TraceIn_ManualMode[18] := BenchUut1.ManualMode;
   TraceIn_SingleStepMode[18] := BenchUut1.SingleStepMode;
   TraceIn_SingleCycleMode[18] := BenchUut1.SingleCycleMode;
   TraceIn_ContinuousMode[18] := BenchUut1.ContinuousMode;
   TraceIn_EmergencyStop[18] := BenchUut1.EmergencyStop;
   TraceIn_Start[18] := BenchUut1.Start;
   TraceIn_DownButton[18] := BenchUut1.DownButton;
   TraceIn_UpButton[18] := BenchUut1.UpButton;
   TraceIn_LeftButton[18] := BenchUut1.LeftButton;
   TraceIn_RightButton[18] := BenchUut1.RightButton;
   TraceIn_GripButton[18] := BenchUut1.GripButton;
   TraceIn_ReleaseButton[18] := BenchUut1.ReleaseButton;
   TraceIn_DownLimitSwitch[18] := BenchUut1.DownLimitSwitch;
   TraceIn_UpLimitSwitch[18] := BenchUut1.UpLimitSwitch;
   TraceIn_LeftLimitSwitch[18] := BenchUut1.LeftLimitSwitch;
   TraceIn_RightLimitSwitch[18] := BenchUut1.RightLimitSwitch;
   TraceIn_GripLimitSwitch[18] := BenchUut1.GripLimitSwitch;
   TraceIn_ReleaseLimitSwitch[18] := BenchUut1.ReleaseLimitSwitch;
   BenchUut1();
   TraceOut_MoveDown[18] := BenchUut1.MoveDown;
   TraceOut_MoveUp[18] := BenchUut1.MoveUp;
   TraceOut_MoveLeft[18] := BenchUut1.MoveLeft;
   TraceOut_MoveRight[18] := BenchUut1.MoveRight;
   TraceOut_ActivateGrip[18] := BenchUut1.ActivateGrip;
   TraceOut_ActivateRelease[18] := BenchUut1.ActivateRelease;
   BenchCalls := BenchCalls + 1;
 19:
   BenchUut2.ManualMode := FALSE;
   BenchUut2.SingleStepMode := FALSE;
   BenchUut2.SingleCycleMode := TRUE;
   BenchUut2.ContinuousMode := FALSE;
   BenchUut2.EmergencyStop := TRUE;
   BenchUut2.Start := FALSE;
   BenchUut2.DownButton := FALSE;
   BenchUut2.UpButton := FALSE;
   BenchUut2.LeftButton := FALSE;
   BenchUut2.RightButton := FALSE;
   BenchUut2.GripButton := FALSE;
   BenchUut2.ReleaseButton := FALSE;
   BenchUut2.DownLimitSwitch := FALSE;
   BenchUut2.UpLimitSwitch := TRUE;
   BenchUut2.LeftLimitSwitch := TRUE;
   BenchUut2.RightLimitSwitch := FALSE;
   BenchUut2.GripLimitSwitch := FALSE;
   BenchUut2.ReleaseLimitSwitch := TRUE;
   TraceIn_ManualMode[19] := BenchUut2.ManualMode;
   TraceIn_SingleStepMode[19] := BenchUut2.SingleStepMode;
   TraceIn_SingleCycleMode[19] := BenchUut2.SingleCycleMode;
   TraceIn_ContinuousMode[19] := BenchUut2.ContinuousMode;
   TraceIn_EmergencyStop[19] := BenchUut2.EmergencyStop;
   TraceIn_Start[19] := BenchUut2.Start;
   TraceIn_DownButton[19] := BenchUut2.DownButton;
   TraceIn_UpButton[19] := BenchUut2.UpButton;
   TraceIn_LeftButton[19] := BenchUut2.LeftButton;
   TraceIn_RightButton[19] := BenchUut2.RightButton;
   TraceIn_GripButton[19] := BenchUut2.GripButton;
   TraceIn_ReleaseButton[19] := BenchUut2.ReleaseButton;
   TraceIn_DownLimitSwitch[19] := BenchUut2.DownLimitSwitch;
   TraceIn_UpLimitSwitch[19] := BenchUut2.UpLimitSwitch;
   TraceIn_LeftLimitSwitch[19] := BenchUut2.LeftLimitSwitch;
   TraceIn_RightLimitSwitch[19] := BenchUut2.RightLimitSwitch;
   TraceIn_GripLimitSwitch[19] := BenchUut2.GripLimitSwitch;
   TraceIn_ReleaseLimitSwitch[19] := BenchUut2.ReleaseLimitSwitch;
   BenchUut2();
   TraceOut_MoveDown[19] := BenchUut2.MoveDown;
   TraceOut_MoveUp[19] := BenchUut2.MoveUp;
   TraceOut_MoveLeft[19] := BenchUut2.MoveLeft;
   TraceOut_MoveRight[19] := BenchUut2.MoveRight;
   TraceOut_ActivateGrip[19] := BenchUut2.ActivateGrip;
   TraceOut_ActivateRelease[19] := BenchUut2.ActivateRelease;
   BenchCalls := BenchCalls + 1;
 20:
   BenchUut2.ManualMode := FALSE;
   BenchUut2.SingleStepMode := FALSE;
   BenchUut2.SingleCycleMode := TRUE;
   BenchUut2.ContinuousMode := FALSE;
   BenchUut2.EmergencyStop := TRUE;
   BenchUut2.Start := TRUE;
   BenchUut2.DownButton := FALSE;
   BenchUut2.UpButton := FALSE;
   BenchUut2.LeftButton := FALSE;
   BenchUut2.RightButton := FALSE;
   BenchUut2.GripButton := FALSE;
   BenchUut2.ReleaseButton := FALSE;
   BenchUut2.DownLimitSwitch := FALSE;
   BenchUut2.UpLimitSwitch := TRUE;
   BenchUut2.LeftLimitSwitch := TRUE;
   BenchUut2.RightLimitSwitch := FALSE;
   BenchUut2.GripLimitSwitch := FALSE;
   BenchUut2.ReleaseLimitSwitch := TRUE;
   TraceIn_ManualMode[20] := BenchUut2.ManualMode;
   TraceIn_SingleStepMode[20] := BenchUut2.SingleStepMode;
   TraceIn_SingleCycleMode[20] := BenchUut2.SingleCycleMode;
   TraceIn_ContinuousMode[20] := BenchUut2.ContinuousMode;
   TraceIn_EmergencyStop[20] := BenchUut2.EmergencyStop;
   TraceIn_Start[20] := BenchUut2.Start;
   TraceIn_DownButton[20] := BenchUut2.DownButton;
   TraceIn_UpButton[20] := BenchUut2.UpButton;
   TraceIn_LeftButton[20] := BenchUut2.LeftButton;
   TraceIn_RightButton[20] := BenchUut2.RightButton;
   TraceIn_GripButton[20] := BenchUut2.GripButton;
   TraceIn_ReleaseButton[20] := BenchUut2.ReleaseButton;
   TraceIn_DownLimitSwitch[20] := BenchUut2.DownLimitSwitch;
   TraceIn_UpLimitSwitch[20] := BenchUut2.UpLimitSwitch;
   TraceIn_LeftLimitSwitch[20] := BenchUut2.LeftLimitSwitch;
   TraceIn_RightLimitSwitch[20] := BenchUut2.RightLimitSwitch;
   TraceIn_GripLimitSwitch[20] := BenchUut2.GripLimitSwitch;
   TraceIn_ReleaseLimitSwitch[20] := BenchUut2.ReleaseLimitSwitch;
   BenchUut2();
   TraceOut_MoveDown[20] := BenchUut2.MoveDown;
   TraceOut_MoveUp[20] := BenchUut2.MoveUp;
   TraceOut_MoveLeft[20] := BenchUut2.MoveLeft;
   TraceOut_MoveRight[20] := BenchUut2.MoveRight;
   TraceOut_ActivateGrip[20] := BenchUut2.ActivateGrip;
   TraceOut_ActivateRelease[20] := BenchUut2.ActivateRelease;
   BenchCalls := BenchCalls + 1;
 21:
   BenchUut2.ManualMode := FALSE;
   BenchUut2.SingleStepMode := FALSE;
   BenchUut2.SingleCycleMode := TRUE;
   BenchUut2.ContinuousMode := FALSE;
   BenchUut2.EmergencyStop := TRUE;
   BenchUut2.Start := FALSE;
   BenchUut2.DownButton := FALSE;
   BenchUut2.UpButton := FALSE;
   BenchUut2.LeftButton := FALSE;
   BenchUut2.RightButton := FALSE;
   BenchUut2.GripButton := FALSE;
   BenchUut2.ReleaseButton := FALSE;
   BenchUut2.DownLimitSwitch := TRUE;
   BenchUut2.UpLimitSwitch := FALSE;
   BenchUut2.LeftLimitSwitch := TRUE;
   BenchUut2.RightLimitSwitch := FALSE;
   BenchUut2.GripLimitSwitch := FALSE;
   BenchUut2.ReleaseLimitSwitch := FALSE;
   TraceIn_ManualMode[21] := BenchUut2.ManualMode;
   TraceIn_SingleStepMode[21] := BenchUut2.SingleStepMode;
   TraceIn_SingleCycleMode[21] := BenchUut2.SingleCycleMode;
   TraceIn_ContinuousMode[21] := BenchUut2.ContinuousMode;
   TraceIn_EmergencyStop[21] := BenchUut2.EmergencyStop;
   TraceIn_Start[21] := BenchUut2.Start;
   TraceIn_DownButton[21] := BenchUut2.DownButton;
   TraceIn_UpButton[21] := BenchUut2.UpButton;
   TraceIn_LeftButton[21] := BenchUut2.LeftButton;
   TraceIn_RightButton[21] := BenchUut2.RightButton;
   TraceIn_GripButton[21] := BenchUut2.GripButton;
   TraceIn_ReleaseButton[21] := BenchUut2.ReleaseButton;
   TraceIn_DownLimitSwitch[21] := BenchUut2.DownLimitSwitch;
   TraceIn_UpLimitSwitch[21] := BenchUut2.UpLimitSwitch;
   TraceIn_LeftLimitSwitch[21] := BenchUut2.LeftLimitSwitch;
   TraceIn_RightLimitSwitch[21] := BenchUut2.RightLimitSwitch;
   TraceIn_GripLimitSwitch[21] := BenchUut2.GripLimitSwitch;
   TraceIn_ReleaseLimitSwitch[21] := BenchUut2.ReleaseLimitSwitch;
   BenchUut2();
   TraceOut_MoveDown[21] := BenchUut2.MoveDown;
   TraceOut_MoveUp[21] := BenchUut2.MoveUp;
   TraceOut_MoveLeft[21] := BenchUut2.MoveLeft;
   TraceOut_MoveRight[21] := BenchUut2.MoveRight;
   TraceOut_ActivateGrip[21] := BenchUut2.ActivateGrip;
   TraceOut_ActivateRelease[21] := BenchUut2.ActivateRelease;
   BenchCalls := BenchCalls + 1;
 22:
   BenchUut2.ManualMode := FALSE;
   BenchUut2.SingleStepMode := FALSE;
   BenchUut2.SingleCycleMode := TRUE;
   BenchUut2.ContinuousMode := FALSE;
   BenchUut2.EmergencyStop := TRUE;
   BenchUut2.Start := FALSE;
   BenchUut2.DownButton := FALSE;
   BenchUut2.UpButton := FALSE;
   BenchUut2.LeftButton := FALSE;
   BenchUut2.RightButton := FALSE;
   BenchUut2.GripButton := FALSE;
   BenchUut2.ReleaseButton := FALSE;
   BenchUut2.DownLimitSwitch := TRUE;
   BenchUut2.UpLimitSwitch := FALSE;
   BenchUut2.LeftLimitSwitch := TRUE;
   BenchUut2.RightLimitSwitch := FALSE;
   BenchUut2.GripLimitSwitch := TRUE;
   BenchUut2.ReleaseLimitSwitch := FALSE;
   TraceIn_ManualMode[22] := BenchUut2.ManualMode;
   TraceIn_SingleStepMode[22] := BenchUut2.SingleStepMode;
   TraceIn_SingleCycleMode[22] := BenchUut2.SingleCycleMode;
   TraceIn_ContinuousMode[22] := BenchUut2.ContinuousMode;
   TraceIn_EmergencyStop[22] := BenchUut2.EmergencyStop;
   TraceIn_Start[22] := BenchUut2.Start;
   TraceIn_DownButton[22] := BenchUut2.DownButton;
   TraceIn_UpButton[22] := BenchUut2.UpButton;
   TraceIn_LeftButton[22] := BenchUut2.LeftButton;
   TraceIn_RightButton[22] := BenchUut2.RightButton;
   TraceIn_GripButton[22] := BenchUut2.GripButton;
   TraceIn_ReleaseButton[22] := BenchUut2.ReleaseButton;
   TraceIn_DownLimitSwitch[22] := BenchUut2.DownLimitSwitch;
   TraceIn_UpLimitSwitch[22] := BenchUut2.UpLimitSwitch;
   TraceIn_LeftLimitSwitch[22] := BenchUut2.LeftLimitSwitch;
   TraceIn_RightLimitSwitch[22] := BenchUut2.RightLimitSwitch;
   TraceIn_GripLimitSwitch[22] := BenchUut2.GripLimitSwitch;
   TraceIn_ReleaseLimitSwitch[22] := BenchUut2.ReleaseLimitSwitch;
   BenchUut2();
   TraceOut_MoveDown[22] := BenchUut2.MoveDown;
   TraceOut_MoveUp[22] := BenchUut2.MoveUp;
   TraceOut_MoveLeft[22] := BenchUut2.MoveLeft;
   TraceOut_MoveRight[22] := BenchUut2.MoveRight;
   TraceOut_ActivateGrip[22] := BenchUut2.ActivateGrip;
   TraceOut_ActivateRelease[22] := BenchUut2.ActivateRelease;
   BenchCalls := BenchCalls + 1;
 23:
   BenchUut2.ManualMode := FALSE;
   BenchUut2.SingleStepMode := FALSE;
   BenchUut2.SingleCycleMode := TRUE;
   BenchUut2.ContinuousMode := FALSE;
   BenchUut2.EmergencyStop := TRUE;
   BenchUut2.Start := FALSE;
   BenchUut2.DownButton := FALSE;
   BenchUut2.UpButton := FALSE;
   BenchUut2.LeftButton := FALSE;
   BenchUut2.RightButton := FALSE;
   BenchUut2.GripButton := FALSE;
   BenchUut2.ReleaseButton := FALSE;
   BenchUut2.DownLimitSwitch := FALSE;
   BenchUut2.UpLimitSwitch := TRUE;
   BenchUut2.LeftLimitSwitch := TRUE;
   BenchUut2.RightLimitSwitch := FALSE;
   BenchUut2.GripLimitSwitch := TRUE;
   BenchUut2.ReleaseLimitSwitch := FALSE;
   TraceIn_ManualMode[23] := BenchUut2.ManualMode;
   TraceIn_SingleStepMode[23] := BenchUut2.SingleStepMode;
   TraceIn_SingleCycleMode[23] := BenchUut2.SingleCycleMode;
   TraceIn_ContinuousMode[23] := BenchUut2.ContinuousMode;
   TraceIn_EmergencyStop[23] := BenchUut2.EmergencyStop;
   TraceIn_Start[23] := BenchUut2.Start;
   TraceIn_DownButton[23] := BenchUut2.DownButton;
   TraceIn_UpButton[23] := BenchUut2.UpButton;
   TraceIn_LeftButton[23] := BenchUut2.LeftButton;
   TraceIn_RightButton[23] := BenchUut2.RightButton;
   TraceIn_GripButton[23] := BenchUut2.GripButton;
   TraceIn_ReleaseButton[23] := BenchUut2.ReleaseButton;
   TraceIn_DownLimitSwitch[23] := BenchUut2.DownLimitSwitch;
   TraceIn_UpLimitSwitch[23] := BenchUut2.UpLimitSwitch;
   TraceIn_LeftLimitSwitch[23] := BenchUut2.LeftLimitSwitch;
   TraceIn_RightLimitSwitch[23] := BenchUut2.RightLimitSwitch;
   TraceIn_GripLimitSwitch[23] := BenchUut2.GripLimitSwitch;
   TraceIn_ReleaseLimitSwitch[23] := BenchUut2.ReleaseLimitSwitch;
   BenchUut2();
   TraceOut_MoveDown[23] := BenchUut2.MoveDown;
   TraceOut_MoveUp[23] := BenchUut2.MoveUp;
   TraceOut_MoveLeft[23] := BenchUut2.MoveLeft;
   TraceOut_MoveRight[23] := BenchUut2.MoveRight;
   TraceOut_ActivateGrip[23] := BenchUut2.ActivateGrip;
   TraceOut_ActivateRelease[23] := BenchUut2.ActivateRelease;
   BenchCalls := BenchCalls + 1;
 24:
   BenchUut2.ManualMode := FALSE;
   BenchUut2.SingleStepMode := FALSE;
   BenchUut2.SingleCycleMode := TRUE;
   BenchUut2.ContinuousMode := FALSE;
   BenchUut2.EmergencyStop := TRUE;
   BenchUut2.Start := FALSE;
   BenchUut2.DownButton := FALSE;
   BenchUut2.UpButton := FALSE;
   BenchUut2.LeftButton := FALSE;
   BenchUut2.RightButton := FALSE;
   BenchUut2.GripButton := FALSE;
   BenchUut2.ReleaseButton := FALSE;
   BenchUut2.DownLimitSwitch := FALSE;
   BenchUut2.UpLimitSwitch := TRUE;
   BenchUut2.LeftLimitSwitch := FALSE;
   BenchUut2.RightLimitSwitch := TRUE;
   BenchUut2.GripLimitSwitch := TRUE;
   BenchUut2.ReleaseLimitSwitch := FALSE;
   TraceIn_ManualMode[24] := BenchUut2.ManualMode;
   TraceIn_SingleStepMode[24] := BenchUut2.SingleStepMode;
   TraceIn_SingleCycleMode[24] := BenchUut2.SingleCycleMode;
   TraceIn_ContinuousMode[24] := BenchUut2.ContinuousMode;
   TraceIn_EmergencyStop[24] := BenchUut2.EmergencyStop;
   TraceIn_Start[24] := BenchUut2.Start;
   TraceIn_DownButton[24] := BenchUut2.DownButton;
   TraceIn_UpButton[24] := BenchUut2.UpButton;
   TraceIn_LeftButton[24] := BenchUut2.LeftButton;
   TraceIn_RightButton[24] := BenchUut2.RightButton;
   TraceIn_GripButton[24] := BenchUut2.GripButton;
   TraceIn_ReleaseButton[24] := BenchUut2.ReleaseButton;
   TraceIn_DownLimitSwitch[24] := BenchUut2.DownLimitSwitch;
   TraceIn_UpLimitSwitch[24] := BenchUut2.UpLimitSwitch;
   TraceIn_LeftLimitSwitch[24] := BenchUut2.LeftLimitSwitch;
   TraceIn_RightLimitSwitch[24] := BenchUut2.RightLimitSwitch;
   TraceIn_GripLimitSwitch[24] := BenchUut2.GripLimitSwitch;
   TraceIn_ReleaseLimitSwitch[24] := BenchUut2.ReleaseLimitSwitch;
   BenchUut2();
   TraceOut_MoveDown[24] := BenchUut2.MoveDown;
   TraceOut_MoveUp[24] := BenchUut2.MoveUp;
   TraceOut_MoveLeft[24] := BenchUut2.MoveLeft;
   TraceOut_MoveRight[24] := BenchUut2.MoveRight;
   TraceOut_ActivateGrip[24] := BenchUut2.ActivateGrip;
   TraceOut_ActivateRelease[24] := BenchUut2.ActivateRelease;
   BenchCalls := BenchCalls + 1;
 25:
   BenchUut2.ManualMode := FALSE;
   BenchUut2.SingleStepMode := FALSE;
   BenchUut2.SingleCycleMode := TRUE;
   BenchUut2.ContinuousMode := FALSE;
   BenchUut2.EmergencyStop := TRUE;
   BenchUut2.Start := FALSE;
   BenchUut2.DownButton := FALSE;
   BenchUut2.UpButton := FALSE;
   BenchUut2.LeftButton := FALSE;
   BenchUut2.RightButton := FALSE;
   BenchUut2.GripButton := FALSE;
   BenchUut2.ReleaseButton := FALSE;
   BenchUut2.DownLimitSwitch := TRUE;
   BenchUut2.UpLimitSwitch := FALSE;
   BenchUut2.LeftLimitSwitch := FALSE;
   BenchUut2.RightLimitSwitch := TRUE;
   BenchUut2.GripLimitSwitch := FALSE;
   BenchUut2.ReleaseLimitSwitch := FALSE;
   TraceIn_ManualMode[25] := BenchUut2.ManualMode;
   TraceIn_SingleStepMode[25] := BenchUut2.SingleStepMode;
   TraceIn_SingleCycleMode[25] := BenchUut2.SingleCycleMode;
   TraceIn_ContinuousMode[25] := BenchUut2.ContinuousMode;
   TraceIn_EmergencyStop[25] := BenchUut2.EmergencyStop;
   TraceIn_Start[25] := BenchUut2.Start;
   TraceIn_DownButton[25] := BenchUut2.DownButton;
   TraceIn_UpButton[25] := BenchUut2.UpButton;
   TraceIn_LeftButton[25] := BenchUut2.LeftButton;
   TraceIn_RightButton[25] := BenchUut2.RightButton;
   TraceIn_GripButton[25] := BenchUut2.GripButton;
   TraceIn_ReleaseButton[25] := BenchUut2.ReleaseButton;
   TraceIn_DownLimitSwitch[25] := BenchUut2.DownLimitSwitch;
   TraceIn_UpLimitSwitch[25] := BenchUut2.UpLimitSwitch;
   TraceIn_LeftLimitSwitch[25] := BenchUut2.LeftLimitSwitch;
   TraceIn_RightLimitSwitch[25] := BenchUut2.RightLimitSwitch;
   TraceIn_GripLimitSwitch[25] := BenchUut2.GripLimitSwitch;
   TraceIn_ReleaseLimitSwitch[25] := BenchUut2.ReleaseLimitSwitch;
   BenchUut2();
   TraceOut_MoveDown[25] := BenchUut2.MoveDown;
   TraceOut_MoveUp[25] := BenchUut2.MoveUp;
   TraceOut_MoveLeft[25] := BenchUut2.MoveLeft;
   TraceOut_MoveRight[25] := BenchUut2.MoveRight;
   TraceOut_ActivateGrip[25] := BenchUut2.ActivateGrip;
   TraceOut_ActivateRelease[25] := BenchUut2.ActivateRelease;
   BenchCalls := BenchCalls + 1;
 26:
   BenchUut2.ManualMode := FALSE;
   BenchUut2.SingleStepMode := FALSE;
   BenchUut2.SingleCycleMode := TRUE;
   BenchUut2.ContinuousMode := FALSE;
   BenchUut2.EmergencyStop := TRUE;
   BenchUut2.Start := FALSE;
   BenchUut2.DownButton := FALSE;
   BenchUut2.UpButton := FALSE;
   BenchUut2.LeftButton := FALSE;
   BenchUut2.RightButton := FALSE;
   BenchUut2.GripButton := FALSE;
   BenchUut2.ReleaseButton := FALSE;
   BenchUut2.DownLimitSwitch := TRUE;
   BenchUut2.UpLimitSwitch := FALSE;
   BenchUut2.LeftLimitSwitch := FALSE;
   BenchUut2.RightLimitSwitch := TRUE;
   BenchUut2.GripLimitSwitch := FALSE;
   BenchUut2.ReleaseLimitSwitch := TRUE;
   TraceIn_ManualMode[26] := BenchUut2.ManualMode;
   TraceIn_SingleStepMode[26] := BenchUut2.SingleStepMode;
   TraceIn_SingleCycleMode[26] := BenchUut2.SingleCycleMode;
   TraceIn_ContinuousMode[26] := BenchUut2.ContinuousMode;
   TraceIn_EmergencyStop[26] := BenchUut2.EmergencyStop;
   TraceIn_Start[26] := BenchUut2.Start;
   TraceIn_DownButton[26] := BenchUut2.DownButton;
   TraceIn_UpButton[26] := BenchUut2.UpButton;
   TraceIn_LeftButton[26] := BenchUut2.LeftButton;
   TraceIn_RightButton[26] := BenchUut2.RightButton;
   TraceIn_GripButton[26] := BenchUut2.GripButton;
   TraceIn_ReleaseButton[26] := BenchUut2.ReleaseButton;
   TraceIn_DownLimitSwitch[26] := BenchUut2.DownLimitSwitch;
   TraceIn_UpLimitSwitch[26] := BenchUut2.UpLimitSwitch;
   TraceIn_LeftLimitSwitch[26] := BenchUut2.LeftLimitSwitch;
   TraceIn_RightLimitSwitch[26] := BenchUut2.RightLimitSwitch;
   TraceIn_GripLimitSwitch[26] := BenchUut2.GripLimitSwitch;
   TraceIn_ReleaseLimitSwitch[26] := BenchUut2.ReleaseLimitSwitch;
   BenchUut2();
   TraceOut_MoveDown[26] := BenchUut2.MoveDown;
   TraceOut_MoveUp[26] := BenchUut2.MoveUp;
   TraceOut_MoveLeft[26] := BenchUut2.MoveLeft;
   TraceOut_MoveRight[26] := BenchUut2.MoveRight;
   TraceOut_ActivateGrip[26] := BenchUut2.ActivateGrip;
   TraceOut_ActivateRelease[26] := BenchUut2.ActivateRelease;
   BenchCalls := BenchCalls + 1;
 27:
   BenchUut2.ManualMode := FALSE;
   BenchUut2.SingleStepMode := FALSE;
   BenchUut2.SingleCycleMode := TRUE;
   BenchUut2.ContinuousMode := FALSE;
   BenchUut2.EmergencyStop := TRUE;
   BenchUut2.Start := FALSE;
   BenchUut2.DownButton := FALSE;
   BenchUut2.UpButton := FALSE;
   BenchUut2.LeftButton := FALSE;
   BenchUut2.RightButton := FALSE;
   BenchUut2.GripButton := FALSE;
   BenchUut2.ReleaseButton := FALSE;
   BenchUut2.DownLimitSwitch := FALSE;
   BenchUut2.UpLimitSwitch := TRUE;
   BenchUut2.LeftLimitSwitch := FALSE;
   BenchUut2.RightLimitSwitch := TRUE;
   BenchUut2.GripLimitSwitch := FALSE;
   BenchUut2.ReleaseLimitSwitch := TRUE;
   TraceIn_ManualMode[27] := BenchUut2.ManualMode;
   TraceIn_SingleStepMode[27] := BenchUut2.SingleStepMode;
   TraceIn_SingleCycleMode[27] := BenchUut2.SingleCycleMode;
   TraceIn_ContinuousMode[27] := BenchUut2.ContinuousMode;
   TraceIn_EmergencyStop[27] := BenchUut2.EmergencyStop;
   TraceIn_Start[27] := BenchUut2.Start;
   TraceIn_DownButton[27] := BenchUut2.DownButton;
   TraceIn_UpButton[27] := BenchUut2.UpButton;
   TraceIn_LeftButton[27] := BenchUut2.LeftButton;
   TraceIn_RightButton[27] := BenchUut2.RightButton;
   TraceIn_GripButton[27] := BenchUut2.GripButton;
   TraceIn_ReleaseButton[27] := BenchUut2.ReleaseButton;
   TraceIn_DownLimitSwitch[27] := BenchUut2.DownLimitSwitch;
   TraceIn_UpLimitSwitch[27] := BenchUut2.UpLimitSwitch;
   TraceIn_LeftLimitSwitch[27] := BenchUut2.LeftLimitSwitch;
   TraceIn_RightLimitSwitch[27] := BenchUut2.RightLimitSwitch;
   TraceIn_GripLimitSwitch[27] := BenchUut2.GripLimitSwitch;
   TraceIn_ReleaseLimitSwitch[27] := BenchUut2.ReleaseLimitSwitch;
   BenchUut2();
   TraceOut_MoveDown[27] := BenchUut2.MoveDown;
   TraceOut_MoveUp[27] := BenchUut2.MoveUp;
   TraceOut_MoveLeft[27] := BenchUut2.MoveLeft;
   TraceOut_MoveRight[27] := BenchUut2.MoveRight;
   TraceOut_ActivateGrip[27] := BenchUut2.ActivateGrip;
   TraceOut_ActivateRelease[27] := BenchUut2.ActivateRelease;
   BenchCalls := BenchCalls + 1;
 28:
   BenchUut2.ManualMode := FALSE;
   BenchUut2.SingleStepMode := FALSE;
   BenchUut2.SingleCycleMode := TRUE;
   BenchUut2.ContinuousMode := FALSE;
   BenchUut2.EmergencyStop := TRUE;
   BenchUut2.Start := FALSE;
   BenchUut2.DownButton := FALSE;
   BenchUut2.UpButton := FALSE;
   BenchUut2.LeftButton := FALSE;
   BenchUut2.RightButton := FALSE;
   BenchUut2.GripButton := FALSE;
   BenchUut2.ReleaseButton := FALSE;
   BenchUut2.DownLimitSwitch := FALSE;
   BenchUut2.UpLimitSwitch := TRUE;
   BenchUut2.LeftLimitSwitch := TRUE;
   BenchUut2.RightLimitSwitch := FALSE;
   BenchUut2.GripLimitSwitch := FALSE;
   BenchUut2.ReleaseLimitSwitch := TRUE;
   TraceIn_ManualMode[28] := BenchUut2.ManualMode;
   TraceIn_SingleStepMode[28] := BenchUut2.SingleStepMode;
   TraceIn_SingleCycleMode[28] := BenchUut2.SingleCycleMode;
   TraceIn_ContinuousMode[28] := BenchUut2.ContinuousMode;
   TraceIn_EmergencyStop[28] := BenchUut2.EmergencyStop;
   TraceIn_Start[28] := BenchUut2.Start;
   TraceIn_DownButton[28] := BenchUut2.DownButton;
   TraceIn_UpButton[28] := BenchUut2.UpButton;
   TraceIn_LeftButton[28] := BenchUut2.LeftButton;
   TraceIn_RightButton[28] := BenchUut2.RightButton;
   TraceIn_GripButton[28] := BenchUut2.GripButton;
   TraceIn_ReleaseButton[28] := BenchUut2.ReleaseButton;
   TraceIn_DownLimitSwitch[28] := BenchUut2.DownLimitSwitch;
   TraceIn_UpLimitSwitch[28] := BenchUut2.UpLimitSwitch;
   TraceIn_LeftLimitSwitch[28] := BenchUut2.LeftLimitSwitch;
   TraceIn_RightLimitSwitch[28] := BenchUut2.RightLimitSwitch;
   TraceIn_GripLimitSwitch[28] := BenchUut2.GripLimitSwitch;
   TraceIn_ReleaseLimitSwitch[28] := BenchUut2.ReleaseLimitSwitch;
   BenchUut2();
   TraceOut_MoveDown[28] := BenchUut2.MoveDown;
   TraceOut_MoveUp[28] := BenchUut2.MoveUp;
   TraceOut_MoveLeft[28] := BenchUut2.MoveLeft;
   TraceOut_MoveRight[28] := BenchUut2.MoveRight;
   TraceOut_ActivateGrip[28] := BenchUut2.ActivateGrip;
   TraceOut_ActivateRelease[28] := BenchUut2.ActivateRelease;
   BenchCalls := BenchCalls + 1;
 29:
   BenchUut3.ManualMode := FALSE;
   BenchUut3.SingleStepMode := FALSE;
   BenchUut3.SingleCycleMode := FALSE;
   BenchUut3.ContinuousMode := TRUE;
   BenchUut3.EmergencyStop := TRUE;
   BenchUut3.Start := FALSE;
   BenchUut3.DownButton := FALSE;
   BenchUut3.UpButton := FALSE;
   BenchUut3.LeftButton := FALSE;
   BenchUut3.RightButton := FALSE;
   BenchUut3.GripButton := FALSE;
   BenchUut3.ReleaseButton := FALSE;
   BenchUut3.DownLimitSwitch := FALSE;
   BenchUut3.UpLimitSwitch := TRUE;
   BenchUut3.LeftLimitSwitch := TRUE;
   BenchUut3.RightLimitSwitch := FALSE;
   BenchUut3.GripLimitSwitch := FALSE;
   BenchUut3.ReleaseLimitSwitch := TRUE;
   TraceIn_ManualMode[29] := BenchUut3.ManualMode;
   TraceIn_SingleStepMode[29] := BenchUut3.SingleStepMode;
   TraceIn_SingleCycleMode[29] := BenchUut3.SingleCycleMode;
   TraceIn_ContinuousMode[29] := BenchUut3.ContinuousMode;
   TraceIn_EmergencyStop[29] := BenchUut3.EmergencyStop;
   TraceIn_Start[29] := BenchUut3.Start;
   TraceIn_DownButton[29] := BenchUut3.DownButton;
   TraceIn_UpButton[29] := BenchUut3.UpButton;
   TraceIn_LeftButton[29] := BenchUut3.LeftButton;
   TraceIn_RightButton[29] := BenchUut3.RightButton;
   TraceIn_GripButton[29] := BenchUut3.GripButton;
   TraceIn_ReleaseButton[29] := BenchUut3.ReleaseButton;
   TraceIn_DownLimitSwitch[29] := BenchUut3.DownLimitSwitch;
   TraceIn_UpLimitSwitch[29] := BenchUut3.UpLimitSwitch;
   TraceIn_LeftLimitSwitch[29] := BenchUut3.LeftLimitSwitch;
   TraceIn_RightLimitSwitch[29] := BenchUut3.RightLimitSwitch;
   TraceIn_GripLimitSwitch[29] := BenchUut3.GripLimitSwitch;
   TraceIn_ReleaseLimitSwitch[29] := BenchUut3.ReleaseLimitSwitch;
   BenchUut3();
   TraceOut_MoveDown[29] := BenchUut3.MoveDown;
   TraceOut_MoveUp[29] := BenchUut3.MoveUp;
   TraceOut_MoveLeft[29] := BenchUut3.MoveLeft;
   TraceOut_MoveRight[29] := BenchUut3.MoveRight;
   TraceOut_ActivateGrip[29] := BenchUut3.ActivateGrip;
   TraceOut_ActivateRelease[29] := BenchUut3.ActivateRelease;
   BenchCalls := BenchCalls + 1;
 30:
   BenchUut3.ManualMode := FALSE;
   BenchUut3.SingleStepMode := FALSE;
   BenchUut3.SingleCycleMode := FALSE;
   BenchUut3.ContinuousMode := TRUE;
   BenchUut3.EmergencyStop := TRUE;
   BenchUut3.Start := TRUE;
   BenchUut3.DownButton := FALSE;
   BenchUut3.UpButton := FALSE;
   BenchUut3.LeftButton := FALSE;
   BenchUut3.RightButton := FALSE;
   BenchUut3.GripButton := FALSE;
   BenchUut3.ReleaseButton := FALSE;
   BenchUut3.DownLimitSwitch := FALSE;
   BenchUut3.UpLimitSwitch := TRUE;
   BenchUut3.LeftLimitSwitch := TRUE;
   BenchUut3.RightLimitSwitch := FALSE;
   BenchUut3.GripLimitSwitch := FALSE;
   BenchUut3.ReleaseLimitSwitch := TRUE;
   TraceIn_ManualMode[30] := BenchUut3.ManualMode;
   TraceIn_SingleStepMode[30] := BenchUut3.SingleStepMode;
   TraceIn_SingleCycleMode[30] := BenchUut3.SingleCycleMode;
   TraceIn_ContinuousMode[30] := BenchUut3.ContinuousMode;
   TraceIn_EmergencyStop[30] := BenchUut3.EmergencyStop;
   TraceIn_Start[30] := BenchUut3.Start;
   TraceIn_DownButton[30] := BenchUut3.DownButton;
   TraceIn_UpButton[30] := BenchUut3.UpButton;
   TraceIn_LeftButton[30] := BenchUut3.LeftButton;
   TraceIn_RightButton[30] := BenchUut3.RightButton;
   TraceIn_GripButton[30] := BenchUut3.GripButton;
   TraceIn_ReleaseButton[30] := BenchUut3.ReleaseButton;
   TraceIn_DownLimitSwitch[30] := BenchUut3.DownLimitSwitch;
   TraceIn_UpLimitSwitch[30] := BenchUut3.UpLimitSwitch;
   TraceIn_LeftLimitSwitch[30] := BenchUut3.LeftLimitSwitch;
   TraceIn_RightLimitSwitch[30] := BenchUut3.RightLimitSwitch;
   TraceIn_GripLimitSwitch[30] := BenchUut3.GripLimitSwitch;
   TraceIn_ReleaseLimitSwitch[30] := BenchUut3.ReleaseLimitSwitch;
   BenchUut3();
   TraceOut_MoveDown[30] := BenchUut3.MoveDown;
   TraceOut_MoveUp[30] := BenchUut3.MoveUp;
   TraceOut_MoveLeft[30] := BenchUut3.MoveLeft;
   TraceOut_MoveRight[30] := BenchUut3.MoveRight;
   TraceOut_ActivateGrip[30] := BenchUut3.ActivateGrip;
   TraceOut_ActivateRelease[30] := BenchUut3.ActivateRelease;
   BenchCalls := BenchCalls + 1;
 31:
   BenchUut3.ManualMode := FALSE;
   BenchUut3.SingleStepMode := FALSE;
   BenchUut3.SingleCycleMode := FALSE;
   BenchUut3.ContinuousMode := TRUE;
   BenchUut3.EmergencyStop := TRUE;
   BenchUut3.Start := FALSE;
   BenchUut3.DownButton := FALSE;
   BenchUut3.UpButton := FALSE;
   BenchUut3.LeftButton := FALSE;
   BenchUut3.RightButton := FALSE;
   BenchUut3.GripButton := FALSE;
   BenchUut3.ReleaseButton := FALSE;
   BenchUut3.DownLimitSwitch := TRUE;
   BenchUut3.UpLimitSwitch := FALSE;
   BenchUut3.LeftLimitSwitch := TRUE;
   BenchUut3.RightLimitSwitch := FALSE;
   BenchUut3.GripLimitSwitch := FALSE;
   BenchUut3.ReleaseLimitSwitch := FALSE;
   TraceIn_ManualMode[31] := BenchUut3.ManualMode;
   TraceIn_SingleStepMode[31] := BenchUut3.SingleStepMode;
   TraceIn_SingleCycleMode[31] := BenchUut3.SingleCycleMode;
   TraceIn_ContinuousMode[31] := BenchUut3.ContinuousMode;
   TraceIn_EmergencyStop[31] := BenchUut3.EmergencyStop;
   TraceIn_Start[31] := BenchUut3.Start;
   TraceIn_DownButton[31] := BenchUut3.DownButton;
   TraceIn_UpButton[31] := BenchUut3.UpButton;
   TraceIn_LeftButton[31] := BenchUut3.LeftButton;
   TraceIn_RightButton[31] := BenchUut3.RightButton;
   TraceIn_GripButton[31] := BenchUut3.GripButton;
   TraceIn_ReleaseButton[31] := BenchUut3.ReleaseButton;
   TraceIn_DownLimitSwitch[31] := BenchUut3.DownLimitSwitch;
   TraceIn_UpLimitSwitch[31] := BenchUut3.UpLimitSwitch;
   TraceIn_LeftLimitSwitch[31] := BenchUut3.LeftLimitSwitch;
   TraceIn_RightLimitSwitch[31] := BenchUut3.RightLimitSwitch;
   TraceIn_GripLimitSwitch[31] := BenchUut3.GripLimitSwitch;
   TraceIn_ReleaseLimitSwitch[31] := BenchUut3.ReleaseLimitSwitch;
   BenchUut3();
   TraceOut_MoveDown[31] := BenchUut3.MoveDown;
   TraceOut_MoveUp[31] := BenchUut3.MoveUp;
   TraceOut_MoveLeft[31] := BenchUut3.MoveLeft;
   TraceOut_MoveRight[31] := BenchUut3.MoveRight;
   TraceOut_ActivateGrip[31] := BenchUut3.ActivateGrip;
   TraceOut_ActivateRelease[31] := BenchUut3.ActivateRelease;
   BenchCalls := BenchCalls + 1;
 32:
   BenchUut3.ManualMode := FALSE;
   BenchUut3.SingleStepMode := FALSE;
   BenchUut3.SingleCycleMode := FALSE;
   BenchUut3.ContinuousMode := TRUE;
   BenchUut3.EmergencyStop := TRUE;
   BenchUut3.Start := FALSE;
   BenchUut3.DownButton := FALSE;
   BenchUut3.UpButton := FALSE;
   BenchUut3.LeftButton := FALSE;
   BenchUut3.RightButton := FALSE;
   BenchUut3.GripButton := FALSE;
   BenchUut3.ReleaseButton := FALSE;
   BenchUut3.DownLimitSwitch := TRUE;
   BenchUut3.UpLimitSwitch := FALSE;
   BenchUut3.LeftLimitSwitch := TRUE;
   BenchUut3.RightLimitSwitch := FALSE;
   BenchUut3.GripLimitSwitch := TRUE;
   BenchUut3.ReleaseLimitSwitch := FALSE;
   TraceIn_ManualMode[32] := BenchUut3.ManualMode;
   TraceIn_SingleStepMode[32] := BenchUut3.SingleStepMode;
   TraceIn_SingleCycleMode[32] := BenchUut3.SingleCycleMode;
   TraceIn_ContinuousMode[32] := BenchUut3.ContinuousMode;
   TraceIn_EmergencyStop[32] := BenchUut3.EmergencyStop;
   TraceIn_Start[32] := BenchUut3.Start;
   TraceIn_DownButton[32] := BenchUut3.DownButton;
   TraceIn_UpButton[32] := BenchUut3.UpButton;
   TraceIn_LeftButton[32] := BenchUut3.LeftButton;
   TraceIn_RightButton[32] := BenchUut3.RightButton;
   TraceIn_GripButton[32] := BenchUut3.GripButton;
   TraceIn_ReleaseButton[32] := BenchUut3.ReleaseButton;
   TraceIn_DownLimitSwitch[32] := BenchUut3.DownLimitSwitch;
   TraceIn_UpLimitSwitch[32] := BenchUut3.UpLimitSwitch;
   TraceIn_LeftLimitSwitch[32] := BenchUut3.LeftLimitSwitch;
   TraceIn_RightLimitSwitch[32] := BenchUut3.RightLimitSwitch;
   TraceIn_GripLimitSwitch[32] := BenchUut3.GripLimitSwitch;
   TraceIn_ReleaseLimitSwitch[32] := BenchUut3.ReleaseLimitSwitch;
   BenchUut3();
   TraceOut_MoveDown[32] := BenchUut3.MoveDown;
   TraceOut_MoveUp[32] := BenchUut3.MoveUp;
   TraceOut_MoveLeft[32] := BenchUut3.MoveLeft;
   TraceOut_MoveRight[32] := BenchUut3.MoveRight;
   TraceOut_ActivateGrip[32] := BenchUut3.ActivateGrip;
   TraceOut_ActivateRelease[32] := BenchUut3.ActivateRelease;
   BenchCalls := BenchCalls + 1;
 33:
   BenchUut3.ManualMode := FALSE;
   BenchUut3.SingleStepMode := FALSE;
   BenchUut3.SingleCycleMode := FALSE;
   BenchUut3.ContinuousMode := TRUE;
   BenchUut3.EmergencyStop := TRUE;
   BenchUut3.Start := FALSE;
   BenchUut3.DownButton := FALSE;
   BenchUut3.UpButton := FALSE;
   BenchUut3.LeftButton := FALSE;
   BenchUut3.RightButton := FALSE;
   BenchUut3.GripButton := FALSE;
   BenchUut3.ReleaseButton := FALSE;
   BenchUut3.DownLimitSwitch := FALSE;
   BenchUut3.UpLimitSwitch := TRUE;
   BenchUut3.LeftLimitSwitch := TRUE;
   BenchUut3.RightLimitSwitch := FALSE;
   BenchUut3.GripLimitSwitch := TRUE;
   BenchUut3.ReleaseLimitSwitch := FALSE;
   TraceIn_ManualMode[33] := BenchUut3.ManualMode;
   TraceIn_SingleStepMode[33] := BenchUut3.SingleStepMode;
   TraceIn_SingleCycleMode[33] := BenchUut3.SingleCycleMode;
   TraceIn_ContinuousMode[33] := BenchUut3.ContinuousMode;
   TraceIn_EmergencyStop[33] := BenchUut3.EmergencyStop;
   TraceIn_Start[33] := BenchUut3.Start;
   TraceIn_DownButton[33] := BenchUut3.DownButton;
   TraceIn_UpButton[33] := BenchUut3.UpButton;
   TraceIn_LeftButton[33] := BenchUut3.LeftButton;
   TraceIn_RightButton[33] := BenchUut3.RightButton;
   TraceIn_GripButton[33] := BenchUut3.GripButton;
   TraceIn_ReleaseButton[33] := BenchUut3.ReleaseButton;
   TraceIn_DownLimitSwitch[33] := BenchUut3.DownLimitSwitch;
   TraceIn_UpLimitSwitch[33] := BenchUut3.UpLimitSwitch;
   TraceIn_LeftLimitSwitch[33] := BenchUut3.LeftLimitSwitch;
   TraceIn_RightLimitSwitch[33] := BenchUut3.RightLimitSwitch;
   TraceIn_GripLimitSwitch[33] := BenchUut3.GripLimitSwitch;
   TraceIn_ReleaseLimitSwitch[33] := BenchUut3.ReleaseLimitSwitch;
   BenchUut3();
   TraceOut_MoveDown[33] := BenchUut3.MoveDown;
   TraceOut_MoveUp[33] := BenchUut3.MoveUp;
   TraceOut_MoveLeft[33] := BenchUut3.MoveLeft;
   TraceOut_MoveRight[33] := BenchUut3.MoveRight;
   TraceOut_ActivateGrip[33] := BenchUut3.ActivateGrip;
   TraceOut_ActivateRelease[33] := BenchUut3.ActivateRelease;
   BenchCalls := BenchCalls + 1;
 34:
   BenchUut3.ManualMode := FALSE;
   BenchUut3.SingleStepMode := FALSE;
   BenchUut3.SingleCycleMode := FALSE;
   BenchUut3.ContinuousMode := TRUE;
   BenchUut3.EmergencyStop := TRUE;
   BenchUut3.Start := FALSE;
   BenchUut3.DownButton := FALSE;
   BenchUut3.UpButton := FALSE;
   BenchUut3.LeftButton := FALSE;
   BenchUut3.RightButton := FALSE;
   BenchUut3.GripButton := FALSE;
   BenchUut3.ReleaseButton := FALSE;
   BenchUut3.DownLimitSwitch := FALSE;
   BenchUut3.UpLimitSwitch := TRUE;
   BenchUut3.LeftLimitSwitch := FALSE;
   BenchUut3.RightLimitSwitch := TRUE;
   BenchUut3.GripLimitSwitch := TRUE;
   BenchUut3.ReleaseLimitSwitch := FALSE;
   TraceIn_ManualMode[34] := BenchUut3.ManualMode;
   TraceIn_SingleStepMode[34] := BenchUut3.SingleStepMode;
   TraceIn_SingleCycleMode[34] := BenchUut3.SingleCycleMode;
   TraceIn_ContinuousMode[34] := BenchUut3.ContinuousMode;
   TraceIn_EmergencyStop[34] := BenchUut3.EmergencyStop;
   TraceIn_Start[34] := BenchUut3.Start;
   TraceIn_DownButton[34] := BenchUut3.DownButton;
   TraceIn_UpButton[34] := BenchUut3.UpButton;
   TraceIn_LeftButton[34] := BenchUut3.LeftButton;
   TraceIn_RightButton[34] := BenchUut3.RightButton;
   TraceIn_GripButton[34] := BenchUut3.GripButton;
   TraceIn_ReleaseButton[34] := BenchUut3.ReleaseButton;
   TraceIn_DownLimitSwitch[34] := BenchUut3.DownLimitSwitch;
   TraceIn_UpLimitSwitch[34] := BenchUut3.UpLimitSwitch;
   TraceIn_LeftLimitSwitch[34] := BenchUut3.LeftLimitSwitch;
   TraceIn_RightLimitSwitch[34] := BenchUut3.RightLimitSwitch;
   TraceIn_GripLimitSwitch[34] := BenchUut3.GripLimitSwitch;
   TraceIn_ReleaseLimitSwitch[34] := BenchUut3.ReleaseLimitSwitch;
   BenchUut3();
   TraceOut_MoveDown[34] := BenchUut3.MoveDown;
   TraceOut_MoveUp[34] := BenchUut3.MoveUp;
   TraceOut_MoveLeft[34] := BenchUut3.MoveLeft;
   TraceOut_MoveRight[34] := BenchUut3.MoveRight;
   TraceOut_ActivateGrip[34] := BenchUut3.ActivateGrip;
   TraceOut_ActivateRelease[34] := BenchUut3.ActivateRelease;
   BenchCalls := BenchCalls + 1;
 35:
   BenchUut3.ManualMode := FALSE;
   BenchUut3.SingleStepMode := FALSE;
   BenchUut3.SingleCycleMode := FALSE;
   BenchUut3.ContinuousMode := TRUE;
   BenchUut3.EmergencyStop := TRUE;
   BenchUut3.Start := FALSE;
   BenchUut3.DownButton := FALSE;
   BenchUut3.UpButton := FALSE;
   BenchUut3.LeftButton := FALSE;
   BenchUut3.RightButton := FALSE;
   BenchUut3.GripButton := FALSE;
   BenchUut3.ReleaseButton := FALSE;
   BenchUut3.DownLimitSwitch := TRUE;
   BenchUut3.UpLimitSwitch := FALSE;
   BenchUut3.LeftLimitSwitch := FALSE;
   BenchUut3.RightLimitSwitch := TRUE;
   BenchUut3.GripLimitSwitch := FALSE;
   BenchUut3.ReleaseLimitSwitch := FALSE;
   TraceIn_ManualMode[35] := BenchUut3.ManualMode;
   TraceIn_SingleStepMode[35] := BenchUut3.SingleStepMode;
   TraceIn_SingleCycleMode[35] := BenchUut3.SingleCycleMode;
   TraceIn_ContinuousMode[35] := BenchUut3.ContinuousMode;
   TraceIn_EmergencyStop[35] := BenchUut3.EmergencyStop;
   TraceIn_Start[35] := BenchUut3.Start;
   TraceIn_DownButton[35] := BenchUut3.DownButton;
   TraceIn_UpButton[35] := BenchUut3.UpButton;
   TraceIn_LeftButton[35] := BenchUut3.LeftButton;
   TraceIn_RightButton[35] := BenchUut3.RightButton;
   TraceIn_GripButton[35] := BenchUut3.GripButton;
   TraceIn_ReleaseButton[35] := BenchUut3.ReleaseButton;
   TraceIn_DownLimitSwitch[35] := BenchUut3.DownLimitSwitch;
   TraceIn_UpLimitSwitch[35] := BenchUut3.UpLimitSwitch;
   TraceIn_LeftLimitSwitch[35] := BenchUut3.LeftLimitSwitch;
   TraceIn_RightLimitSwitch[35] := BenchUut3.RightLimitSwitch;
   TraceIn_GripLimitSwitch[35] := BenchUut3.GripLimitSwitch;
   TraceIn_ReleaseLimitSwitch[35] := BenchUut3.ReleaseLimitSwitch;
   BenchUut3();
   TraceOut_MoveDown[35] := BenchUut3.MoveDown;
   TraceOut_MoveUp[35] := BenchUut3.MoveUp;
   TraceOut_MoveLeft[35] := BenchUut3.MoveLeft;
   TraceOut_MoveRight[35] := BenchUut3.MoveRight;
   TraceOut_ActivateGrip[35] := BenchUut3.ActivateGrip;
   TraceOut_ActivateRelease[35] := BenchUut3.ActivateRelease;
   BenchCalls := BenchCalls + 1;
 36:
   BenchUut3.ManualMode := FALSE;
   BenchUut3.SingleStepMode := FALSE;
   BenchUut3.SingleCycleMode := FALSE;
   BenchUut3.ContinuousMode := TRUE;
   BenchUut3.EmergencyStop := TRUE;
   BenchUut3.Start := FALSE;
   BenchUut3.DownButton := FALSE;
   BenchUut3.UpButton := FALSE;
   BenchUut3.LeftButton := FALSE;
   BenchUut3.RightButton := FALSE;
   BenchUut3.GripButton := FALSE;
   BenchUut3.ReleaseButton := FALSE;
   BenchUut3.DownLimitSwitch := TRUE;
   BenchUut3.UpLimitSwitch := FALSE;
   BenchUut3.LeftLimitSwitch := FALSE;
   BenchUut3.RightLimitSwitch := TRUE;
   BenchUut3.GripLimitSwitch := FALSE;
   BenchUut3.ReleaseLimitSwitch := TRUE;
   TraceIn_ManualMode[36] := BenchUut3.ManualMode;
   TraceIn_SingleStepMode[36] := BenchUut3.SingleStepMode;
   TraceIn_SingleCycleMode[36] := BenchUut3.SingleCycleMode;
   TraceIn_ContinuousMode[36] := BenchUut3.ContinuousMode;
   TraceIn_EmergencyStop[36] := BenchUut3.EmergencyStop;
   TraceIn_Start[36] := BenchUut3.Start;
   TraceIn_DownButton[36] := BenchUut3.DownButton;
   TraceIn_UpButton[36] := BenchUut3.UpButton;
   TraceIn_LeftButton[36] := BenchUut3.LeftButton;
   TraceIn_RightButton[36] := BenchUut3.RightButton;
   TraceIn_GripButton[36] := BenchUut3.GripButton;
   TraceIn_ReleaseButton[36] := BenchUut3.ReleaseButton;
   TraceIn_DownLimitSwitch[36] := BenchUut3.DownLimitSwitch;
   TraceIn_UpLimitSwitch[36] := BenchUut3.UpLimitSwitch;
   TraceIn_LeftLimitSwitch[36] := BenchUut3.LeftLimitSwitch;
   TraceIn_RightLimitSwitch[36] := BenchUut3.RightLimitSwitch;
   TraceIn_GripLimitSwitch[36] := BenchUut3.GripLimitSwitch;
   TraceIn_ReleaseLimitSwitch[36] := BenchUut3.ReleaseLimitSwitch;
   BenchUut3();
   TraceOut_MoveDown[36] := BenchUut3.MoveDown;
   TraceOut_MoveUp[36] := BenchUut3.MoveUp;
   TraceOut_MoveLeft[36] := BenchUut3.MoveLeft;
   TraceOut_MoveRight[36] := BenchUut3.MoveRight;
   TraceOut_ActivateGrip[36] := BenchUut3.ActivateGrip;
   TraceOut_ActivateRelease[36] := BenchUut3.ActivateRelease;
   BenchCalls := BenchCalls + 1;
 37:
   BenchUut3.ManualMode := FALSE;
   BenchUut3.SingleStepMode := FALSE;
   BenchUut3.SingleCycleMode := FALSE;
   BenchUut3.ContinuousMode := TRUE;
   BenchUut3.EmergencyStop := TRUE;
   BenchUut3.Start := FALSE;
   BenchUut3.DownButton := FALSE;
   BenchUut3.UpButton := FALSE;
   BenchUut3.LeftButton := FALSE;
   BenchUut3.RightButton := FALSE;
   BenchUut3.GripButton := FALSE;
   BenchUut3.ReleaseButton := FALSE;
   BenchUut3.DownLimitSwitch := FALSE;
   BenchUut3.UpLimitSwitch := TRUE;
   BenchUut3.LeftLimitSwitch := FALSE;
   BenchUut3.RightLimitSwitch := TRUE;
   BenchUut3.GripLimitSwitch := FALSE;
   BenchUut3.ReleaseLimitSwitch := TRUE;
   TraceIn_ManualMode[37] := BenchUut3.ManualMode;
   TraceIn_SingleStepMode[37] := BenchUut3.SingleStepMode;
   TraceIn_SingleCycleMode[37] := BenchUut3.SingleCycleMode;
   TraceIn_ContinuousMode[37] := BenchUut3.ContinuousMode;
   TraceIn_EmergencyStop[37] := BenchUut3.EmergencyStop;
   TraceIn_Start[37] := BenchUut3.Start;
   TraceIn_DownButton[37] := BenchUut3.DownButton;
   TraceIn_UpButton[37] := BenchUut3.UpButton;
   TraceIn_LeftButton[37] := BenchUut3.LeftButton;
   TraceIn_RightButton[37] := BenchUut3.RightButton;
   TraceIn_GripButton[37] := BenchUut3.GripButton;
   TraceIn_ReleaseButton[37] := BenchUut3.ReleaseButton;
   TraceIn_DownLimitSwitch[37] := BenchUut3.DownLimitSwitch;
   TraceIn_UpLimitSwitch[37] := BenchUut3.UpLimitSwitch;
   TraceIn_LeftLimitSwitch[37] := BenchUut3.LeftLimitSwitch;
   TraceIn_RightLimitSwitch[37] := BenchUut3.RightLimitSwitch;
   TraceIn_GripLimitSwitch[37] := BenchUut3.GripLimitSwitch;
   TraceIn_ReleaseLimitSwitch[37] := BenchUut3.ReleaseLimitSwitch;
   BenchUut3();
   TraceOut_MoveDown[37] := BenchUut3.MoveDown;
   TraceOut_MoveUp[37] := BenchUut3.MoveUp;
   TraceOut_MoveLeft[37] := BenchUut3.MoveLeft;
   TraceOut_MoveRight[37] := BenchUut3.MoveRight;
   TraceOut_ActivateGrip[37] := BenchUut3.ActivateGrip;
   TraceOut_ActivateRelease[37] := BenchUut3.ActivateRelease;
   BenchCalls := BenchCalls + 1;
 38:
   BenchUut3.ManualMode := FALSE;
   BenchUut3.SingleStepMode := FALSE;
   BenchUut3.SingleCycleMode := FALSE;
   BenchUut3.ContinuousMode := TRUE;
   BenchUut3.EmergencyStop := TRUE;
   BenchUut3.Start := FALSE;
   BenchUut3.DownButton := FALSE;
   BenchUut3.UpButton := FALSE;
   BenchUut3.LeftButton := FALSE;
   BenchUut3.RightButton := FALSE;
   BenchUut3.GripButton := FALSE;
   BenchUut3.ReleaseButton := FALSE;
   BenchUut3.DownLimitSwitch := FALSE;
   BenchUut3.UpLimitSwitch := TRUE;
   BenchUut3.LeftLimitSwitch := TRUE;
   BenchUut3.RightLimitSwitch := FALSE;
   BenchUut3.GripLimitSwitch := FALSE;
   BenchUut3.ReleaseLimitSwitch := TRUE;
   TraceIn_ManualMode[38] := BenchUut3.ManualMode;
   TraceIn_SingleStepMode[38] := BenchUut3.SingleStepMode;
   TraceIn_SingleCycleMode[38] := BenchUut3.SingleCycleMode;
   TraceIn_ContinuousMode[38] := BenchUut3.ContinuousMode;
   TraceIn_EmergencyStop[38] := BenchUut3.EmergencyStop;
   TraceIn_Start[38] := BenchUut3.Start;
   TraceIn_DownButton[38] := BenchUut3.DownButton;
   TraceIn_UpButton[38] := BenchUut3.UpButton;
   TraceIn_LeftButton[38] := BenchUut3.LeftButton;
   TraceIn_RightButton[38] := BenchUut3.RightButton;
   TraceIn_GripButton[38] := BenchUut3.GripButton;
   TraceIn_ReleaseButton[38] := BenchUut3.ReleaseButton;
   TraceIn_DownLimitSwitch[38] := BenchUut3.DownLimitSwitch;
   TraceIn_UpLimitSwitch[38] := BenchUut3.UpLimitSwitch;
   TraceIn_LeftLimitSwitch[38] := BenchUut3.LeftLimitSwitch;
   TraceIn_RightLimitSwitch[38] := BenchUut3.RightLimitSwitch;
   TraceIn_GripLimitSwitch[38] := BenchUut3.GripLimitSwitch;
   TraceIn_ReleaseLimitSwitch[38] := BenchUut3.ReleaseLimitSwitch;
   BenchUut3();
   TraceOut_MoveDown[38] := BenchUut3.MoveDown;
   TraceOut_MoveUp[38] := BenchUut3.MoveUp;
   TraceOut_MoveLeft[38] := BenchUut3.MoveLeft;
   TraceOut_MoveRight[38] := BenchUut3.MoveRight;
   TraceOut_ActivateGrip[38] := BenchUut3.ActivateGrip;
   TraceOut_ActivateRelease[38] := BenchUut3.ActivateRelease;
   BenchCalls := BenchCalls + 1;
 39:
   BenchUut4.ManualMode := FALSE;
   BenchUut4.SingleStepMode := FALSE;
   BenchUut4.SingleCycleMode := TRUE;
   BenchUut4.ContinuousMode := FALSE;
   BenchUut4.EmergencyStop := TRUE;
   BenchUut4.Start := FALSE;
   BenchUut4.DownButton := FALSE;
   BenchUut4.UpButton := FALSE;
   BenchUut4.LeftButton := FALSE;
   BenchUut4.RightButton := FALSE;
   BenchUut4.GripButton := FALSE;
   BenchUut4.ReleaseButton := FALSE;
   BenchUut4.DownLimitSwitch := FALSE;
   BenchUut4.UpLimitSwitch := TRUE;
   BenchUut4.LeftLimitSwitch := TRUE;
   BenchUut4.RightLimitSwitch := FALSE;
   BenchUut4.GripLimitSwitch := FALSE;
   BenchUut4.ReleaseLimitSwitch := TRUE;
   TraceIn_ManualMode[39] := BenchUut4.ManualMode;
   TraceIn_SingleStepMode[39] := BenchUut4.SingleStepMode;
   TraceIn_SingleCycleMode[39] := BenchUut4.SingleCycleMode;
   TraceIn_ContinuousMode[39] := BenchUut4.ContinuousMode;
   TraceIn_EmergencyStop[39] := BenchUut4.EmergencyStop;
   TraceIn_Start[39] := BenchUut4.Start;
   TraceIn_DownButton[39] := BenchUut4.DownButton;
   TraceIn_UpButton[39] := BenchUut4.UpButton;
   TraceIn_LeftButton[39] := BenchUut4.LeftButton;
   TraceIn_RightButton[39] := BenchUut4.RightButton;
   TraceIn_GripButton[39] := BenchUut4.GripButton;
   TraceIn_ReleaseButton[39] := BenchUut4.ReleaseButton;
   TraceIn_DownLimitSwitch[39] := BenchUut4.DownLimitSwitch;
   TraceIn_UpLimitSwitch[39] := BenchUut4.UpLimitSwitch;
   TraceIn_LeftLimitSwitch[39] := BenchUut4.LeftLimitSwitch;
   TraceIn_RightLimitSwitch[39] := BenchUut4.RightLimitSwitch;
   TraceIn_GripLimitSwitch[39] := BenchUut4.GripLimitSwitch;
   TraceIn_ReleaseLimitSwitch[39] := BenchUut4.ReleaseLimitSwitch;
   BenchUut4();
   TraceOut_MoveDown[39] := BenchUut4.MoveDown;
   TraceOut_MoveUp[39] := BenchUut4.MoveUp;
   TraceOut_MoveLeft[39] := BenchUut4.MoveLeft;
   TraceOut_MoveRight[39] := BenchUut4.MoveRight;
   TraceOut_ActivateGrip[39] := BenchUut4.ActivateGrip;
   TraceOut_ActivateRelease[39] := BenchUut4.ActivateRelease;
   BenchCalls := BenchCalls + 1;
 40:
   BenchUut4.ManualMode := FALSE;
   BenchUut4.SingleStepMode := FALSE;
   BenchUut4.SingleCycleMode := TRUE;
   BenchUut4.ContinuousMode := FALSE;
   BenchUut4.EmergencyStop := TRUE;
   BenchUut4.Start := TRUE;
   BenchUut4.DownButton := FALSE;
   BenchUut4.UpButton := FALSE;
   BenchUut4.LeftButton := FALSE;
   BenchUut4.RightButton := FALSE;
   BenchUut4.GripButton := FALSE;
   BenchUut4.ReleaseButton := FALSE;
   BenchUut4.DownLimitSwitch := FALSE;
   BenchUut4.UpLimitSwitch := TRUE;
   BenchUut4.LeftLimitSwitch := TRUE;
   BenchUut4.RightLimitSwitch := FALSE;
   BenchUut4.GripLimitSwitch := FALSE;
   BenchUut4.ReleaseLimitSwitch := TRUE;
   TraceIn_ManualMode[40] := BenchUut4.ManualMode;
   TraceIn_SingleStepMode[40] := BenchUut4.SingleStepMode;
   TraceIn_SingleCycleMode[40] := BenchUut4.SingleCycleMode;
   TraceIn_ContinuousMode[40] := BenchUut4.ContinuousMode;
   TraceIn_EmergencyStop[40] := BenchUut4.EmergencyStop;
   TraceIn_Start[40] := BenchUut4.Start;
   TraceIn_DownButton[40] := BenchUut4.DownButton;
   TraceIn_UpButton[40] := BenchUut4.UpButton;
   TraceIn_LeftButton[40] := BenchUut4.LeftButton;
   TraceIn_RightButton[40] := BenchUut4.RightButton;
   TraceIn_GripButton[40] := BenchUut4.GripButton;
   TraceIn_ReleaseButton[40] := BenchUut4.ReleaseButton;
   TraceIn_DownLimitSwitch[40] := BenchUut4.DownLimitSwitch;
   TraceIn_UpLimitSwitch[40] := BenchUut4.UpLimitSwitch;
   TraceIn_LeftLimitSwitch[40] := BenchUut4.LeftLimitSwitch;
   TraceIn_RightLimitSwitch[40] := BenchUut4.RightLimitSwitch;
   TraceIn_GripLimitSwitch[40] := BenchUut4.GripLimitSwitch;
   TraceIn_ReleaseLimitSwitch[40] := BenchUut4.ReleaseLimitSwitch;
   BenchUut4();
   TraceOut_MoveDown[40] := BenchUut4.MoveDown;
   TraceOut_MoveUp[40] := BenchUut4.MoveUp;
   TraceOut_MoveLeft[40] := BenchUut4.MoveLeft;
   TraceOut_MoveRight[40] := BenchUut4.MoveRight;
   TraceOut_ActivateGrip[40] := BenchUut4.ActivateGrip;
   TraceOut_ActivateRelease[40] := BenchUut4.ActivateRelease;
   BenchCalls := BenchCalls + 1;
 41:
   BenchUut4.ManualMode := FALSE;
   BenchUut4.SingleStepMode := FALSE;
   BenchUut4.SingleCycleMode := TRUE;
   BenchUut4.ContinuousMode := FALSE;
   BenchUut4.EmergencyStop := FALSE;
   BenchUut4.Start := FALSE;
   BenchUut4.DownButton := FALSE;
   BenchUut4.UpButton := FALSE;
   BenchUut4.LeftButton := FALSE;
   BenchUut4.RightButton := FALSE;
   BenchUut4.GripButton := FALSE;
   BenchUut4.ReleaseButton := FALSE;
   BenchUut4.DownLimitSwitch := FALSE;
   BenchUut4.UpLimitSwitch := FALSE;
   BenchUut4.LeftLimitSwitch := TRUE;
   BenchUut4.RightLimitSwitch := FALSE;
   BenchUut4.GripLimitSwitch := FALSE;
   BenchUut4.ReleaseLimitSwitch := TRUE;
   TraceIn_ManualMode[41] := BenchUut4.ManualMode;
   TraceIn_SingleStepMode[41] := BenchUut4.SingleStepMode;
   TraceIn_SingleCycleMode[41] := BenchUut4.SingleCycleMode;
   TraceIn_ContinuousMode[41] := BenchUut4.ContinuousMode;
   TraceIn_EmergencyStop[41] := BenchUut4.EmergencyStop;
   TraceIn_Start[41] := BenchUut4.Start;
   TraceIn_DownButton[41] := BenchUut4.DownButton;
   TraceIn_UpButton[41] := BenchUut4.UpButton;
   TraceIn_LeftButton[41] := BenchUut4.LeftButton;
   TraceIn_RightButton[41] := BenchUut4.RightButton;
   TraceIn_GripButton[41] := BenchUut4.GripButton;
   TraceIn_ReleaseButton[41] := BenchUut4.ReleaseButton;
   TraceIn_DownLimitSwitch[41] := BenchUut4.DownLimitSwitch;
   TraceIn_UpLimitSwitch[41] := BenchUut4.UpLimitSwitch;
   TraceIn_LeftLimitSwitch[41] := BenchUut4.LeftLimitSwitch;
   TraceIn_RightLimitSwitch[41] := BenchUut4.RightLimitSwitch;
   TraceIn_GripLimitSwitch[41] := BenchUut4.GripLimitSwitch;
   TraceIn_ReleaseLimitSwitch[41] := BenchUut4.ReleaseLimitSwitch;
   BenchUut4();
   TraceOut_MoveDown[41] := BenchUut4.MoveDown;
   TraceOut_MoveUp[41] := BenchUut4.MoveUp;
   TraceOut_MoveLeft[41] := BenchUut4.MoveLeft;
   TraceOut_MoveRight[41] := BenchUut4.MoveRight;
   TraceOut_ActivateGrip[41] := BenchUut4.ActivateGrip;
   TraceOut_ActivateRelease[41] := BenchUut4.ActivateRelease;
   BenchCalls := BenchCalls + 1;
 42:
   BenchUut4.ManualMode := FALSE;
   BenchUut4.SingleStepMode := FALSE;
   BenchUut4.SingleCycleMode := TRUE;
   BenchUut4.ContinuousMode := FALSE;
   BenchUut4.EmergencyStop := TRUE;
   BenchUut4.Start := FALSE;
   BenchUut4.DownButton := FALSE;
   BenchUut4.UpButton := FALSE;
   BenchUut4.LeftButton := FALSE;
   BenchUut4.RightButton := FALSE;
   BenchUut4.GripButton := FALSE;
   BenchUut4.ReleaseButton := FALSE;
   BenchUut4.DownLimitSwitch := FALSE;
   BenchUut4.UpLimitSwitch := FALSE;
   BenchUut4.LeftLimitSwitch := TRUE;
   BenchUut4.RightLimitSwitch := FALSE;
   BenchUut4.GripLimitSwitch := FALSE;
   BenchUut4.ReleaseLimitSwitch := TRUE;
   TraceIn_ManualMode[42] := BenchUut4.ManualMode;
   TraceIn_SingleStepMode[42] := BenchUut4.SingleStepMode;
   TraceIn_SingleCycleMode[42] := BenchUut4.SingleCycleMode;
   TraceIn_ContinuousMode[42] := BenchUut4.ContinuousMode;
   TraceIn_EmergencyStop[42] := BenchUut4.EmergencyStop;
   TraceIn_Start[42] := BenchUut4.Start;
   TraceIn_DownButton[42] := BenchUut4.DownButton;
   TraceIn_UpButton[42] := BenchUut4.UpButton;
   TraceIn_LeftButton[42] := BenchUut4.LeftButton;
   TraceIn_RightButton[42] := BenchUut4.RightButton;
   TraceIn_GripButton[42] := BenchUut4.GripButton;
   TraceIn_ReleaseButton[42] := BenchUut4.ReleaseButton;
   TraceIn_DownLimitSwitch[42] := BenchUut4.DownLimitSwitch;
   TraceIn_UpLimitSwitch[42] := BenchUut4.UpLimitSwitch;
   TraceIn_LeftLimitSwitch[42] := BenchUut4.LeftLimitSwitch;
   TraceIn_RightLimitSwitch[42] := BenchUut4.RightLimitSwitch;
   TraceIn_GripLimitSwitch[42] := BenchUut4.GripLimitSwitch;
   TraceIn_ReleaseLimitSwitch[42] := BenchUut4.ReleaseLimitSwitch;
   BenchUut4();
   TraceOut_MoveDown[42] := BenchUut4.MoveDown;
   TraceOut_MoveUp[42] := BenchUut4.MoveUp;
   TraceOut_MoveLeft[42] := BenchUut4.MoveLeft;
   TraceOut_MoveRight[42] := BenchUut4.MoveRight;
   TraceOut_ActivateGrip[42] := BenchUut4.ActivateGrip;
   TraceOut_ActivateRelease[42] := BenchUut4.ActivateRelease;
   BenchCalls := BenchCalls + 1;
 43:
   BenchUut4.ManualMode := FALSE;
   BenchUut4.SingleStepMode := FALSE;
   BenchUut4.SingleCycleMode := TRUE;
   BenchUut4.ContinuousMode := FALSE;
   BenchUut4.EmergencyStop := TRUE;
   BenchUut4.Start := FALSE;
   BenchUut4.DownButton := FALSE;
   BenchUut4.UpButton := FALSE;
   BenchUut4.LeftButton := FALSE;
   BenchUut4.RightButton := FALSE;
   BenchUut4.GripButton := FALSE;
   BenchUut4.ReleaseButton := FALSE;
   BenchUut4.DownLimitSwitch := FALSE;
   BenchUut4.UpLimitSwitch := TRUE;
   BenchUut4.LeftLimitSwitch := TRUE;
   BenchUut4.RightLimitSwitch := FALSE;
   BenchUut4.GripLimitSwitch := FALSE;
   BenchUut4.ReleaseLimitSwitch := TRUE;
   TraceIn_ManualMode[43] := BenchUut4.ManualMode;
   TraceIn_SingleStepMode[43] := BenchUut4.SingleStepMode;
   TraceIn_SingleCycleMode[43] := BenchUut4.SingleCycleMode;
   TraceIn_ContinuousMode[43] := BenchUut4.ContinuousMode;
   TraceIn_EmergencyStop[43] := BenchUut4.EmergencyStop;
   TraceIn_Start[43] := BenchUut4.Start;
   TraceIn_DownButton[43] := BenchUut4.DownButton;
   TraceIn_UpButton[43] := BenchUut4.UpButton;
   TraceIn_LeftButton[43] := BenchUut4.LeftButton;
   TraceIn_RightButton[43] := BenchUut4.RightButton;
   TraceIn_GripButton[43] := BenchUut4.GripButton;
   TraceIn_ReleaseButton[43] := BenchUut4.ReleaseButton;
   TraceIn_DownLimitSwitch[43] := BenchUut4.DownLimitSwitch;
   TraceIn_UpLimitSwitch[43] := BenchUut4.UpLimitSwitch;
   TraceIn_LeftLimitSwitch[43] := BenchUut4.LeftLimitSwitch;
   TraceIn_RightLimitSwitch[43] := BenchUut4.RightLimitSwitch;
   TraceIn_GripLimitSwitch[43] := BenchUut4.GripLimitSwitch;
   TraceIn_ReleaseLimitSwitch[43] := BenchUut4.ReleaseLimitSwitch;
   BenchUut4();
   TraceOut_MoveDown[43] := BenchUut4.MoveDown;
   TraceOut_MoveUp[43] := BenchUut4.MoveUp;
   TraceOut_MoveLeft[43] := BenchUut4.MoveLeft;
   TraceOut_MoveRight[43] := BenchUut4.MoveRight;
   TraceOut_ActivateGrip[43] := BenchUut4.ActivateGrip;
   TraceOut_ActivateRelease[43] := BenchUut4.ActivateRelease;
   BenchCalls := BenchCalls + 1;
 44:
   BenchUut4.ManualMode := FALSE;
   BenchUut4.SingleStepMode := FALSE;
   BenchUut4.SingleCycleMode := TRUE;
   BenchUut4.ContinuousMode := FALSE;
   BenchUut4.EmergencyStop := TRUE;
   BenchUut4.Start := TRUE;
   BenchUut4.DownButton := FALSE;
   BenchUut4.UpButton := FALSE;
   BenchUut4.LeftButton := FALSE;
   BenchUut4.RightButton := FALSE;
   BenchUut4.GripButton := FALSE;
   BenchUut4.ReleaseButton := FALSE;
   BenchUut4.DownLimitSwitch := FALSE;
   BenchUut4.UpLimitSwitch := TRUE;
   BenchUut4.LeftLimitSwitch := TRUE;
   BenchUut4.RightLimitSwitch := FALSE;
   BenchUut4.GripLimitSwitch := FALSE;
   BenchUut4.ReleaseLimitSwitch := TRUE;
   TraceIn_ManualMode[44] := BenchUut4.ManualMode;
   TraceIn_SingleStepMode[44] := BenchUut4.SingleStepMode;
   TraceIn_SingleCycleMode[44] := BenchUut4.SingleCycleMode;
   TraceIn_ContinuousMode[44] := BenchUut4.ContinuousMode;
   TraceIn_EmergencyStop[44] := BenchUut4.EmergencyStop;
   TraceIn_Start[44] := BenchUut4.Start;
   TraceIn_DownButton[44] := BenchUut4.DownButton;
   TraceIn_UpButton[44] := BenchUut4.UpButton;
   TraceIn_LeftButton[44] := BenchUut4.LeftButton;
   TraceIn_RightButton[44] := BenchUut4.RightButton;
   TraceIn_GripButton[44] := BenchUut4.GripButton;
   TraceIn_ReleaseButton[44] := BenchUut4.ReleaseButton;
   TraceIn_DownLimitSwitch[44] := BenchUut4.DownLimitSwitch;
   TraceIn_UpLimitSwitch[44] := BenchUut4.UpLimitSwitch;
   TraceIn_LeftLimitSwitch[44] := BenchUut4.LeftLimitSwitch;
   TraceIn_RightLimitSwitch[44] := BenchUut4.RightLimitSwitch;
   TraceIn_GripLimitSwitch[44] := BenchUut4.GripLimitSwitch;
   TraceIn_ReleaseLimitSwitch[44] := BenchUut4.ReleaseLimitSwitch;
   BenchUut4();
   TraceOut_MoveDown[44] := BenchUut4.MoveDown;
   TraceOut_MoveUp[44] := BenchUut4.MoveUp;
   TraceOut_MoveLeft[44] := BenchUut4.MoveLeft;
   TraceOut_MoveRight[44] := BenchUut4.MoveRight;
   TraceOut_ActivateGrip[44] := BenchUut4.ActivateGrip;
   TraceOut_ActivateRelease[44] := BenchUut4.ActivateRelease;
   BenchCalls := BenchCalls + 1;
 45:
   BenchUut5.ManualMode := FALSE;
   BenchUut5.SingleStepMode := FALSE;
   BenchUut5.SingleCycleMode := FALSE;
   BenchUut5.ContinuousMode := FALSE;
   BenchUut5.EmergencyStop := TRUE;
   BenchUut5.Start := FALSE;
   BenchUut5.DownButton := FALSE;
   BenchUut5.UpButton := FALSE;
   BenchUut5.LeftButton := FALSE;
   BenchUut5.RightButton := FALSE;
   BenchUut5.GripButton := FALSE;
   BenchUut5.ReleaseButton := FALSE;
   BenchUut5.DownLimitSwitch := FALSE;
   BenchUut5.UpLimitSwitch := FALSE;
   BenchUut5.LeftLimitSwitch := FALSE;
   BenchUut5.RightLimitSwitch := FALSE;
   BenchUut5.GripLimitSwitch := FALSE;
   BenchUut5.ReleaseLimitSwitch := FALSE;
   TraceIn_ManualMode[45] := BenchUut5.ManualMode;
   TraceIn_SingleStepMode[45] := BenchUut5.SingleStepMode;
   TraceIn_SingleCycleMode[45] := BenchUut5.SingleCycleMode;
   TraceIn_ContinuousMode[45] := BenchUut5.ContinuousMode;
   TraceIn_EmergencyStop[45] := BenchUut5.EmergencyStop;
   TraceIn_Start[45] := BenchUut5.Start;
   TraceIn_DownButton[45] := BenchUut5.DownButton;
   TraceIn_UpButton[45] := BenchUut5.UpButton;
   TraceIn_LeftButton[45] := BenchUut5.LeftButton;
   TraceIn_RightButton[45] := BenchUut5.RightButton;
   TraceIn_GripButton[45] := BenchUut5.GripButton;
   TraceIn_ReleaseButton[45] := BenchUut5.ReleaseButton;
   TraceIn_DownLimitSwitch[45] := BenchUut5.DownLimitSwitch;
   TraceIn_UpLimitSwitch[45] := BenchUut5.UpLimitSwitch;
   TraceIn_LeftLimitSwitch[45] := BenchUut5.LeftLimitSwitch;
   TraceIn_RightLimitSwitch[45] := BenchUut5.RightLimitSwitch;
   TraceIn_GripLimitSwitch[45] := BenchUut5.GripLimitSwitch;
   TraceIn_ReleaseLimitSwitch[45] := BenchUut5.ReleaseLimitSwitch;
   BenchUut5();
   TraceOut_MoveDown[45] := BenchUut5.MoveDown;
   TraceOut_MoveUp[45] := BenchUut5.MoveUp;
   TraceOut_MoveLeft[45] := BenchUut5.MoveLeft;
   TraceOut_MoveRight[45] := BenchUut5.MoveRight;
   TraceOut_ActivateGrip[45] := BenchUut5.ActivateGrip;
   TraceOut_ActivateRelease[45] := BenchUut5.ActivateRelease;
   BenchCalls := BenchCalls + 1;
 46:
   BenchUut5.ManualMode := TRUE;
   BenchUut5.SingleStepMode := FALSE;
   BenchUut5.SingleCycleMode := FALSE;
   BenchUut5.ContinuousMode := FALSE;
   BenchUut5.EmergencyStop := TRUE;
   BenchUut5.Start := FALSE;
   BenchUut5.DownButton := FALSE;
   BenchUut5.UpButton := TRUE;
   BenchUut5.LeftButton := FALSE;
   BenchUut5.RightButton := FALSE;
   BenchUut5.GripButton := TRUE;
   BenchUut5.ReleaseButton := TRUE;
   BenchUut5.DownLimitSwitch := FALSE;
   BenchUut5.UpLimitSwitch := FALSE;
   BenchUut5.LeftLimitSwitch := FALSE;
   BenchUut5.RightLimitSwitch := FALSE;
   BenchUut5.GripLimitSwitch := FALSE;
   BenchUut5.ReleaseLimitSwitch := FALSE;
   TraceIn_ManualMode[46] := BenchUut5.ManualMode;
   TraceIn_SingleStepMode[46] := BenchUut5.SingleStepMode;
   TraceIn_SingleCycleMode[46] := BenchUut5.SingleCycleMode;
   TraceIn_ContinuousMode[46] := BenchUut5.ContinuousMode;
   TraceIn_EmergencyStop[46] := BenchUut5.EmergencyStop;
   TraceIn_Start[46] := BenchUut5.Start;
   TraceIn_DownButton[46] := BenchUut5.DownButton;
   TraceIn_UpButton[46] := BenchUut5.UpButton;
   TraceIn_LeftButton[46] := BenchUut5.LeftButton;
   TraceIn_RightButton[46] := BenchUut5.RightButton;
   TraceIn_GripButton[46] := BenchUut5.GripButton;
   TraceIn_ReleaseButton[46] := BenchUut5.ReleaseButton;
   TraceIn_DownLimitSwitch[46] := BenchUut5.DownLimitSwitch;
   TraceIn_UpLimitSwitch[46] := BenchUut5.UpLimitSwitch;
   TraceIn_LeftLimitSwitch[46] := BenchUut5.LeftLimitSwitch;
   TraceIn_RightLimitSwitch[46] := BenchUut5.RightLimitSwitch;
   TraceIn_GripLimitSwitch[46] := BenchUut5.GripLimitSwitch;
   TraceIn_ReleaseLimitSwitch[46] := BenchUut5.ReleaseLimitSwitch;
   BenchUut5();
   TraceOut_MoveDown[46] := BenchUut5.MoveDown;
   TraceOut_MoveUp[46] := BenchUut5.MoveUp;
   TraceOut_MoveLeft[46] := BenchUut5.MoveLeft;
   TraceOut_MoveRight[46] := BenchUut5.MoveRight;
   TraceOut_ActivateGrip[46] := BenchUut5.ActivateGrip;
   TraceOut_ActivateRelease[46] := BenchUut5.ActivateRelease;
   BenchCalls := BenchCalls + 1;
 47:
   BenchUut5.ManualMode := TRUE;
   BenchUut5.SingleStepMode := FALSE;
   BenchUut5.SingleCycleMode := FALSE;
   BenchUut5.ContinuousMode := FALSE;
   BenchUut5.EmergencyStop := TRUE;
   BenchUut5.Start := FALSE;
   BenchUut5.DownButton := FALSE;
   BenchUut5.UpButton := FALSE;
   BenchUut5.LeftButton := TRUE;
   BenchUut5.RightButton := FALSE;
   BenchUut5.GripButton := FALSE;
   BenchUut5.ReleaseButton := TRUE;
   BenchUut5.DownLimitSwitch := FALSE;
   BenchUut5.UpLimitSwitch := FALSE;
   BenchUut5.LeftLimitSwitch := FALSE;
   BenchUut5.RightLimitSwitch := FALSE;
   BenchUut5.GripLimitSwitch := FALSE;
   BenchUut5.ReleaseLimitSwitch := FALSE;
   TraceIn_ManualMode[47] := BenchUut5.ManualMode;
   TraceIn_SingleStepMode[47] := BenchUut5.SingleStepMode;
   TraceIn_SingleCycleMode[47] := BenchUut5.SingleCycleMode;
   TraceIn_ContinuousMode[47] := BenchUut5.ContinuousMode;
   TraceIn_EmergencyStop[47] := BenchUut5.EmergencyStop;
   TraceIn_Start[47] := BenchUut5.Start;
   TraceIn_DownButton[47] := BenchUut5.DownButton;
   TraceIn_UpButton[47] := BenchUut5.UpButton;
   TraceIn_LeftButton[47] := BenchUut5.LeftButton;
   TraceIn_RightButton[47] := BenchUut5.RightButton;
   TraceIn_GripButton[47] := BenchUut5.GripButton;
   TraceIn_ReleaseButton[47] := BenchUut5.ReleaseButton;
   TraceIn_DownLimitSwitch[47] := BenchUut5.DownLimitSwitch;
   TraceIn_UpLimitSwitch[47] := BenchUut5.UpLimitSwitch;
   TraceIn_LeftLimitSwitch[47] := BenchUut5.LeftLimitSwitch;
   TraceIn_RightLimitSwitch[47] := BenchUut5.RightLimitSwitch;
   TraceIn_GripLimitSwitch[47] := BenchUut5.GripLimitSwitch;
   TraceIn_ReleaseLimitSwitch[47] := BenchUut5.ReleaseLimitSwitch;
   BenchUut5();
   TraceOut_MoveDown[47] := BenchUut5.MoveDown;
   TraceOut_MoveUp[47] := BenchUut5.MoveUp;
   TraceOut_MoveLeft[47] := BenchUut5.MoveLeft;
   TraceOut_MoveRight[47] := BenchUut5.MoveRight;
   TraceOut_ActivateGrip[47] := BenchUut5.ActivateGrip;
   TraceOut_ActivateRelease[47] := BenchUut5.ActivateRelease;
   BenchCalls := BenchCalls + 1;
 48:
   BenchUut5.ManualMode := FALSE;
   BenchUut5.SingleStepMode := TRUE;
   BenchUut5.SingleCycleMode := FALSE;
   BenchUut5.ContinuousMode := FALSE;
   BenchUut5.EmergencyStop := TRUE;
   BenchUut5.Start := TRUE;
   BenchUut5.DownButton := FALSE;
   BenchUut5.UpButton := FALSE;
   BenchUut5.LeftButton := FALSE;
   BenchUut5.RightButton := FALSE;
   BenchUut5.GripButton := FALSE;
   BenchUut5.ReleaseButton := FALSE;
   BenchUut5.DownLimitSwitch := FALSE;
   BenchUut5.UpLimitSwitch := TRUE;
   BenchUut5.LeftLimitSwitch := FALSE;
   BenchUut5.RightLimitSwitch := FALSE;
   BenchUut5.GripLimitSwitch := FALSE;
   BenchUut5.ReleaseLimitSwitch := FALSE;
   TraceIn_ManualMode[48] := BenchUut5.ManualMode;
   TraceIn_SingleStepMode[48] := BenchUut5.SingleStepMode;
   TraceIn_SingleCycleMode[48] := BenchUut5.SingleCycleMode;
   TraceIn_ContinuousMode[48] := BenchUut5.ContinuousMode;
   TraceIn_EmergencyStop[48] := BenchUut5.EmergencyStop;
   TraceIn_Start[48] := BenchUut5.Start;
   TraceIn_DownButton[48] := BenchUut5.DownButton;
   TraceIn_UpButton[48] := BenchUut5.UpButton;
   TraceIn_LeftButton[48] := BenchUut5.LeftButton;
   TraceIn_RightButton[48] := BenchUut5.RightButton;
   TraceIn_GripButton[48] := BenchUut5.GripButton;
   TraceIn_ReleaseButton[48] := BenchUut5.ReleaseButton;
   TraceIn_DownLimitSwitch[48] := BenchUut5.DownLimitSwitch;
   TraceIn_UpLimitSwitch[48] := BenchUut5.UpLimitSwitch;
   TraceIn_LeftLimitSwitch[48] := BenchUut5.LeftLimitSwitch;
   TraceIn_RightLimitSwitch[48] := BenchUut5.RightLimitSwitch;
   TraceIn_GripLimitSwitch[48] := BenchUut5.GripLimitSwitch;
   TraceIn_ReleaseLimitSwitch[48] := BenchUut5.ReleaseLimitSwitch;
   BenchUut5();
   TraceOut_MoveDown[48] := BenchUut5.MoveDown;
   TraceOut_MoveUp[48] := BenchUut5.MoveUp;
   TraceOut_MoveLeft[48] := BenchUut5.MoveLeft;
   TraceOut_MoveRight[48] := BenchUut5.MoveRight;
   TraceOut_ActivateGrip[48] := BenchUut5.ActivateGrip;
   TraceOut_ActivateRelease[48] := BenchUut5.ActivateRelease;
   BenchCalls := BenchCalls + 1;
 49:
   BenchUut5.ManualMode := FALSE;
   BenchUut5.SingleStepMode := TRUE;
   BenchUut5.SingleCycleMode := FALSE;
   BenchUut5.ContinuousMode := FALSE;
   BenchUut5.EmergencyStop := TRUE;
   BenchUut5.Start := TRUE;
   BenchUut5.DownButton := FALSE;
   BenchUut5.UpButton := FALSE;
   BenchUut5.LeftButton := FALSE;
   BenchUut5.RightButton := FALSE;
   BenchUut5.GripButton := FALSE;
   BenchUut5.ReleaseButton := FALSE;
   BenchUut5.DownLimitSwitch := FALSE;
   BenchUut5.UpLimitSwitch := TRUE;
   BenchUut5.LeftLimitSwitch := FALSE;
   BenchUut5.RightLimitSwitch := FALSE;
   BenchUut5.GripLimitSwitch := FALSE;
   BenchUut5.ReleaseLimitSwitch := FALSE;
   TraceIn_ManualMode[49] := BenchUut5.ManualMode;
   TraceIn_SingleStepMode[49] := BenchUut5.SingleStepMode;
   TraceIn_SingleCycleMode[49] := BenchUut5.SingleCycleMode;
   TraceIn_ContinuousMode[49] := BenchUut5.ContinuousMode;
   TraceIn_EmergencyStop[49] := BenchUut5.EmergencyStop;
   TraceIn_Start[49] := BenchUut5.Start;
   TraceIn_DownButton[49] := BenchUut5.DownButton;
   TraceIn_UpButton[49] := BenchUut5.UpButton;
   TraceIn_LeftButton[49] := BenchUut5.LeftButton;
   TraceIn_RightButton[49] := BenchUut5.RightButton;
   TraceIn_GripButton[49] := BenchUut5.GripButton;
   TraceIn_ReleaseButton[49] := BenchUut5.ReleaseButton;
   TraceIn_DownLimitSwitch[49] := BenchUut5.DownLimitSwitch;
   TraceIn_UpLimitSwitch[49] := BenchUut5.UpLimitSwitch;
   TraceIn_LeftLimitSwitch[49] := BenchUut5.LeftLimitSwitch;
   TraceIn_RightLimitSwitch[49] := BenchUut5.RightLimitSwitch;
   TraceIn_GripLimitSwitch[49] := BenchUut5.GripLimitSwitch;
   TraceIn_ReleaseLimitSwitch[49] := BenchUut5.ReleaseLimitSwitch;
   BenchUut5();
   TraceOut_MoveDown[49] := BenchUut5.MoveDown;
   TraceOut_MoveUp[49] := BenchUut5.MoveUp;
   TraceOut_MoveLeft[49] := BenchUut5.MoveLeft;
   TraceOut_MoveRight[49] := BenchUut5.MoveRight;
   TraceOut_ActivateGrip[49] := BenchUut5.ActivateGrip;
   TraceOut_ActivateRelease[49] := BenchUut5.ActivateRelease;
   BenchCalls := BenchCalls + 1;
 50:
   BenchUut5.ManualMode := FALSE;
   BenchUut5.SingleStepMode := TRUE;
   BenchUut5.SingleCycleMode := FALSE;
   BenchUut5.ContinuousMode := FALSE;
   BenchUut5.EmergencyStop := TRUE;
   BenchUut5.Start := FALSE;
   BenchUut5.DownButton := FALSE;
   BenchUut5.UpButton := FALSE;
   BenchUut5.LeftButton := FALSE;
   BenchUut5.RightButton := FALSE;
   BenchUut5.GripButton := FALSE;
   BenchUut5.ReleaseButton := FALSE;
   BenchUut5.DownLimitSwitch := FALSE;
   BenchUut5.UpLimitSwitch := TRUE;
   BenchUut5.LeftLimitSwitch := TRUE;
   BenchUut5.RightLimitSwitch := FALSE;
   BenchUut5.GripLimitSwitch := FALSE;
   BenchUut5.ReleaseLimitSwitch := FALSE;
   TraceIn_ManualMode[50] := BenchUut5.ManualMode;
   TraceIn_SingleStepMode[50] := BenchUut5.SingleStepMode;
   TraceIn_SingleCycleMode[50] := BenchUut5.SingleCycleMode;
   TraceIn_ContinuousMode[50] := BenchUut5.ContinuousMode;
   TraceIn_EmergencyStop[50] := BenchUut5.EmergencyStop;
   TraceIn_Start[50] := BenchUut5.Start;
   TraceIn_DownButton[50] := BenchUut5.DownButton;
   TraceIn_UpButton[50] := BenchUut5.UpButton;
   TraceIn_LeftButton[50] := BenchUut5.LeftButton;
   TraceIn_RightButton[50] := BenchUut5.RightButton;
   TraceIn_GripButton[50] := BenchUut5.GripButton;
   TraceIn_ReleaseButton[50] := BenchUut5.ReleaseButton;
   TraceIn_DownLimitSwitch[50] := BenchUut5.DownLimitSwitch;
   TraceIn_UpLimitSwitch[50] := BenchUut5.UpLimitSwitch;
   TraceIn_LeftLimitSwitch[50] := BenchUut5.LeftLimitSwitch;
   TraceIn_RightLimitSwitch[50] := BenchUut5.RightLimitSwitch;
   TraceIn_GripLimitSwitch[50] := BenchUut5.GripLimitSwitch;
   TraceIn_ReleaseLimitSwitch[50] := BenchUut5.ReleaseLimitSwitch;
   BenchUut5();
   TraceOut_MoveDown[50] := BenchUut5.MoveDown;
   TraceOut_MoveUp[50] := BenchUut5.MoveUp;
   TraceOut_MoveLeft[50] := BenchUut5.MoveLeft;
   TraceOut_MoveRight[50] := BenchUut5.MoveRight;
   TraceOut_ActivateGrip[50] := BenchUut5.ActivateGrip;
   TraceOut_ActivateRelease[50] := BenchUut5.ActivateRelease;
   BenchCalls := BenchCalls + 1;
 51:
   BenchUut5.ManualMode := FALSE;
   BenchUut5.SingleStepMode := TRUE;
   BenchUut5.SingleCycleMode := FALSE;
   BenchUut5.ContinuousMode := FALSE;
   BenchUut5.EmergencyStop := TRUE;
   BenchUut5.Start := TRUE;
   BenchUut5.DownButton := FALSE;
   BenchUut5.UpButton := FALSE;
   BenchUut5.LeftButton := FALSE;
   BenchUut5.RightButton := FALSE;
   BenchUut5.GripButton := FALSE;
   BenchUut5.ReleaseButton := FALSE;
   BenchUut5.DownLimitSwitch := FALSE;
   BenchUut5.UpLimitSwitch := TRUE;
   BenchUut5.LeftLimitSwitch := TRUE;
   BenchUut5.RightLimitSwitch := FALSE;
   BenchUut5.GripLimitSwitch := FALSE;
   BenchUut5.ReleaseLimitSwitch := FALSE;
   TraceIn_ManualMode[51] := BenchUut5.ManualMode;
   TraceIn_SingleStepMode[51] := BenchUut5.SingleStepMode;
   TraceIn_SingleCycleMode[51] := BenchUut5.SingleCycleMode;
   TraceIn_ContinuousMode[51] := BenchUut5.ContinuousMode;
   TraceIn_EmergencyStop[51] := BenchUut5.EmergencyStop;
   TraceIn_Start[51] := BenchUut5.Start;
   TraceIn_DownButton[51] := BenchUut5.DownButton;
   TraceIn_UpButton[51] := BenchUut5.UpButton;
   TraceIn_LeftButton[51] := BenchUut5.LeftButton;
   TraceIn_RightButton[51] := BenchUut5.RightButton;
   TraceIn_GripButton[51] := BenchUut5.GripButton;
   TraceIn_ReleaseButton[51] := BenchUut5.ReleaseButton;
   TraceIn_DownLimitSwitch[51] := BenchUut5.DownLimitSwitch;
   TraceIn_UpLimitSwitch[51] := BenchUut5.UpLimitSwitch;
   TraceIn_LeftLimitSwitch[51] := BenchUut5.LeftLimitSwitch;
   TraceIn_RightLimitSwitch[51] := BenchUut5.RightLimitSwitch;
   TraceIn_GripLimitSwitch[51] := BenchUut5.GripLimitSwitch;
   TraceIn_ReleaseLimitSwitch[51] := BenchUut5.ReleaseLimitSwitch;
   BenchUut5();
   TraceOut_MoveDown[51] := BenchUut5.MoveDown;
   TraceOut_MoveUp[51] := BenchUut5.MoveUp;
   TraceOut_MoveLeft[51] := BenchUut5.MoveLeft;
   TraceOut_MoveRight[51] := BenchUut5.MoveRight;
   TraceOut_ActivateGrip[51] := BenchUut5.ActivateGrip;
   TraceOut_ActivateRelease[51] := BenchUut5.ActivateRelease;
   BenchCalls := BenchCalls + 1;
 52:
   BenchUut5.ManualMode := FALSE;
   BenchUut5.SingleStepMode := TRUE;
   BenchUut5.SingleCycleMode := FALSE;
   BenchUut5.ContinuousMode := FALSE;
   BenchUut5.EmergencyStop := TRUE;
   BenchUut5.Start := FALSE;
   BenchUut5.DownButton := FALSE;
   BenchUut5.UpButton := FALSE;
   BenchUut5.LeftButton := FALSE;
   BenchUut5.RightButton := FALSE;
   BenchUut5.GripButton := FALSE;
   BenchUut5.ReleaseButton := FALSE;
   BenchUut5.DownLimitSwitch := TRUE;
   BenchUut5.UpLimitSwitch := FALSE;
   BenchUut5.LeftLimitSwitch := FALSE;
   BenchUut5.RightLimitSwitch := FALSE;
   BenchUut5.GripLimitSwitch := FALSE;
   BenchUut5.ReleaseLimitSwitch := FALSE;
   TraceIn_ManualMode[52] := BenchUut5.ManualMode;
   TraceIn_SingleStepMode[52] := BenchUut5.SingleStepMode;
   TraceIn_SingleCycleMode[52] := BenchUut5.SingleCycleMode;
   TraceIn_ContinuousMode[52] := BenchUut5.ContinuousMode;
   TraceIn_EmergencyStop[52] := BenchUut5.EmergencyStop;
   TraceIn_Start[52] := BenchUut5.Start;
   TraceIn_DownButton[52] := BenchUut5.DownButton;
   TraceIn_UpButton[52] := BenchUut5.UpButton;
   TraceIn_LeftButton[52] := BenchUut5.LeftButton;
   TraceIn_RightButton[52] := BenchUut5.RightButton;
   TraceIn_GripButton[52] := BenchUut5.GripButton;
   TraceIn_ReleaseButton[52] := BenchUut5.ReleaseButton;
   TraceIn_DownLimitSwitch[52] := BenchUut5.DownLimitSwitch;
   TraceIn_UpLimitSwitch[52] := BenchUut5.UpLimitSwitch;
   TraceIn_LeftLimitSwitch[52] := BenchUut5.LeftLimitSwitch;
   TraceIn_RightLimitSwitch[52] := BenchUut5.RightLimitSwitch;
   TraceIn_GripLimitSwitch[52] := BenchUut5.GripLimitSwitch;
   TraceIn_ReleaseLimitSwitch[52] := BenchUut5.ReleaseLimitSwitch;
   BenchUut5();
   TraceOut_MoveDown[52] := BenchUut5.MoveDown;
   TraceOut_MoveUp[52] := BenchUut5.MoveUp;
   TraceOut_MoveLeft[52] := BenchUut5.MoveLeft;
   TraceOut_MoveRight[52] := BenchUut5.MoveRight;
   TraceOut_ActivateGrip[52] := BenchUut5.ActivateGrip;
   TraceOut_ActivateRelease[52] := BenchUut5.ActivateRelease;
   BenchCalls := BenchCalls + 1;
 53:
   BenchUut5.ManualMode := FALSE;
   BenchUut5.SingleStepMode := TRUE;
   BenchUut5.SingleCycleMode := FALSE;
   BenchUut5.ContinuousMode := FALSE;
   BenchUut5.EmergencyStop := TRUE;
   BenchUut5.Start := TRUE;
   BenchUut5.DownButton := FALSE;
   BenchUut5.UpButton := FALSE;
   BenchUut5.LeftButton := FALSE;
   BenchUut5.RightButton := FALSE;
   BenchUut5.GripButton := FALSE;
   BenchUut5.ReleaseButton := FALSE;
   BenchUut5.DownLimitSwitch := FALSE;
   BenchUut5.UpLimitSwitch := FALSE;
   BenchUut5.LeftLimitSwitch := FALSE;
   BenchUut5.RightLimitSwitch := FALSE;
   BenchUut5.GripLimitSwitch := FALSE;
   BenchUut5.ReleaseLimitSwitch := FALSE;
   TraceIn_ManualMode[53] := BenchUut5.ManualMode;
   TraceIn_SingleStepMode[53] := BenchUut5.SingleStepMode;
   TraceIn_SingleCycleMode[53] := BenchUut5.SingleCycleMode;
   TraceIn_ContinuousMode[53] := BenchUut5.ContinuousMode;
   TraceIn_EmergencyStop[53] := BenchUut5.EmergencyStop;
   TraceIn_Start[53] := BenchUut5.Start;
   TraceIn_DownButton[53] := BenchUut5.DownButton;
   TraceIn_UpButton[53] := BenchUut5.UpButton;
   TraceIn_LeftButton[53] := BenchUut5.LeftButton;
   TraceIn_RightButton[53] := BenchUut5.RightButton;
   TraceIn_GripButton[53] := BenchUut5.GripButton;
   TraceIn_ReleaseButton[53] := BenchUut5.ReleaseButton;
   TraceIn_DownLimitSwitch[53] := BenchUut5.DownLimitSwitch;
   TraceIn_UpLimitSwitch[53] := BenchUut5.UpLimitSwitch;
   TraceIn_LeftLimitSwitch[53] := BenchUut5.LeftLimitSwitch;
   TraceIn_RightLimitSwitch[53] := BenchUut5.RightLimitSwitch;
   TraceIn_GripLimitSwitch[53] := BenchUut5.GripLimitSwitch;
   TraceIn_ReleaseLimitSwitch[53] := BenchUut5.ReleaseLimitSwitch;
   BenchUut5();
   TraceOut_MoveDown[53] := BenchUut5.MoveDown;
   TraceOut_MoveUp[53] := BenchUut5.MoveUp;
   TraceOut_MoveLeft[53] := BenchUut5.MoveLeft;
   TraceOut_MoveRight[53] := BenchUut5.MoveRight;
   TraceOut_ActivateGrip[53] := BenchUut5.ActivateGrip;
   TraceOut_ActivateRelease[53] := BenchUut5.ActivateRelease;
   BenchCalls := BenchCalls + 1;
 54:
   BenchUut5.ManualMode := FALSE;
   BenchUut5.SingleStepMode := TRUE;
   BenchUut5.SingleCycleMode := FALSE;
   BenchUut5.ContinuousMode := FALSE;
   BenchUut5.EmergencyStop := TRUE;
   BenchUut5.Start := FALSE;
   BenchUut5.DownButton := FALSE;
   BenchUut5.UpButton := FALSE;
   BenchUut5.LeftButton := FALSE;
   BenchUut5.RightButton := FALSE;
   BenchUut5.GripButton := FALSE;
   BenchUut5.ReleaseButton := FALSE;
   BenchUut5.DownLimitSwitch := FALSE;
   BenchUut5.UpLimitSwitch := FALSE;
   BenchUut5.LeftLimitSwitch := FALSE;
   BenchUut5.RightLimitSwitch := FALSE;
   BenchUut5.GripLimitSwitch := TRUE;
   BenchUut5.ReleaseLimitSwitch := FALSE;
   TraceIn_ManualMode[54] := BenchUut5.ManualMode;
   TraceIn_SingleStepMode[54] := BenchUut5.SingleStepMode;
   TraceIn_SingleCycleMode[54] := BenchUut5.SingleCycleMode;
   TraceIn_ContinuousMode[54] := BenchUut5.ContinuousMode;
   TraceIn_EmergencyStop[54] := BenchUut5.EmergencyStop;
   TraceIn_Start[54] := BenchUut5.Start;
   TraceIn_DownButton[54] := BenchUut5.DownButton;
   TraceIn_UpButton[54] := BenchUut5.UpButton;
   TraceIn_LeftButton[54] := BenchUut5.LeftButton;
   TraceIn_RightButton[54] := BenchUut5.RightButton;
   TraceIn_GripButton[54] := BenchUut5.GripButton;
   TraceIn_ReleaseButton[54] := BenchUut5.ReleaseButton;
   TraceIn_DownLimitSwitch[54] := BenchUut5.DownLimitSwitch;
   TraceIn_UpLimitSwitch[54] := BenchUut5.UpLimitSwitch;
   TraceIn_LeftLimitSwitch[54] := BenchUut5.LeftLimitSwitch;
   TraceIn_RightLimitSwitch[54] := BenchUut5.RightLimitSwitch;
   TraceIn_GripLimitSwitch[54] := BenchUut5.GripLimitSwitch;
   TraceIn_ReleaseLimitSwitch[54] := BenchUut5.ReleaseLimitSwitch;
   BenchUut5();
   TraceOut_MoveDown[54] := BenchUut5.MoveDown;
   TraceOut_MoveUp[54] := BenchUut5.MoveUp;
   TraceOut_MoveLeft[54] := BenchUut5.MoveLeft;
   TraceOut_MoveRight[54] := BenchUut5.MoveRight;
   TraceOut_ActivateGrip[54] := BenchUut5.ActivateGrip;
   TraceOut_ActivateRelease[54] := BenchUut5.ActivateRelease;
   BenchCalls := BenchCalls + 1;
 55:
   BenchUut5.ManualMode := FALSE;
   BenchUut5.SingleStepMode := TRUE;
   BenchUut5.SingleCycleMode := FALSE;
   BenchUut5.ContinuousMode := FALSE;
   BenchUut5.EmergencyStop := TRUE;
   BenchUut5.Start := TRUE;
   BenchUut5.DownButton := FALSE;
   BenchUut5.UpButton := FALSE;
   BenchUut5.LeftButton := FALSE;
   BenchUut5.RightButton := FALSE;
   BenchUut5.GripButton := FALSE;
   BenchUut5.ReleaseButton := FALSE;
   BenchUut5.DownLimitSwitch := FALSE;
   BenchUut5.UpLimitSwitch := FALSE;
   BenchUut5.LeftLimitSwitch := FALSE;
   BenchUut5.RightLimitSwitch := FALSE;
   BenchUut5.GripLimitSwitch := FALSE;
   BenchUut5.ReleaseLimitSwitch := FALSE;
   TraceIn_ManualMode[55] := BenchUut5.ManualMode;
   TraceIn_SingleStepMode[55] := BenchUut5.SingleStepMode;
   TraceIn_SingleCycleMode[55] := BenchUut5.SingleCycleMode;
   TraceIn_ContinuousMode[55] := BenchUut5.ContinuousMode;
   TraceIn_EmergencyStop[55] := BenchUut5.EmergencyStop;
   TraceIn_Start[55] := BenchUut5.Start;
   TraceIn_DownButton[55] := BenchUut5.DownButton;
   TraceIn_UpButton[55] := BenchUut5.UpButton;
   TraceIn_LeftButton[55] := BenchUut5.LeftButton;
   TraceIn_RightButton[55] := BenchUut5.RightButton;
   TraceIn_GripButton[55] := BenchUut5.GripButton;
   TraceIn_ReleaseButton[55] := BenchUut5.ReleaseButton;
   TraceIn_DownLimitSwitch[55] := BenchUut5.DownLimitSwitch;
   TraceIn_UpLimitSwitch[55] := BenchUut5.UpLimitSwitch;
   TraceIn_LeftLimitSwitch[55] := BenchUut5.LeftLimitSwitch;
   TraceIn_RightLimitSwitch[55] := BenchUut5.RightLimitSwitch;
   TraceIn_GripLimitSwitch[55] := BenchUut5.GripLimitSwitch;
   TraceIn_ReleaseLimitSwitch[55] := BenchUut5.ReleaseLimitSwitch;
   BenchUut5();
   TraceOut_MoveDown[55] := BenchUut5.MoveDown;
   TraceOut_MoveUp[55] := BenchUut5.MoveUp;
   TraceOut_MoveLeft[55] := BenchUut5.MoveLeft;
   TraceOut_MoveRight[55] := BenchUut5.MoveRight;
   TraceOut_ActivateGrip[55] := BenchUut5.ActivateGrip;
   TraceOut_ActivateRelease[55] := BenchUut5.ActivateRelease;
   BenchCalls := BenchCalls + 1;
 56:
   BenchUut5.ManualMode := FALSE;
   BenchUut5.SingleStepMode := TRUE;
   BenchUut5.SingleCycleMode := FALSE;
   BenchUut5.ContinuousMode := FALSE;
   BenchUut5.EmergencyStop := TRUE;
   BenchUut5.Start := FALSE;
   BenchUut5.DownButton := FALSE;
   BenchUut5.UpButton := FALSE;
   BenchUut5.LeftButton := FALSE;
   BenchUut5.RightButton := FALSE;
   BenchUut5.GripButton := FALSE;
   BenchUut5.ReleaseButton := FALSE;
   BenchUut5.DownLimitSwitch := FALSE;
   BenchUut5.UpLimitSwitch := TRUE;
   BenchUut5.LeftLimitSwitch := FALSE;
   BenchUut5.RightLimitSwitch := FALSE;
   BenchUut5.GripLimitSwitch := FALSE;
   BenchUut5.ReleaseLimitSwitch := FALSE;
   TraceIn_ManualMode[56] := BenchUut5.ManualMode;
   TraceIn_SingleStepMode[56] := BenchUut5.SingleStepMode;
   TraceIn_SingleCycleMode[56] := BenchUut5.SingleCycleMode;
   TraceIn_ContinuousMode[56] := BenchUut5.ContinuousMode;
   TraceIn_EmergencyStop[56] := BenchUut5.EmergencyStop;
   TraceIn_Start[56] := BenchUut5.Start;
   TraceIn_DownButton[56] := BenchUut5.DownButton;
   TraceIn_UpButton[56] := BenchUut5.UpButton;
   TraceIn_LeftButton[56] := BenchUut5.LeftButton;
   TraceIn_RightButton[56] := BenchUut5.RightButton;
   TraceIn_GripButton[56] := BenchUut5.GripButton;
   TraceIn_ReleaseButton[56] := BenchUut5.ReleaseButton;
   TraceIn_DownLimitSwitch[56] := BenchUut5.DownLimitSwitch;
   TraceIn_UpLimitSwitch[56] := BenchUut5.UpLimitSwitch;
   TraceIn_LeftLimitSwitch[56] := BenchUut5.LeftLimitSwitch;
   TraceIn_RightLimitSwitch[56] := BenchUut5.RightLimitSwitch;
   TraceIn_GripLimitSwitch[56] := BenchUut5.GripLimitSwitch;
   TraceIn_ReleaseLimitSwitch[56] := BenchUut5.ReleaseLimitSwitch;
   BenchUut5();
   TraceOut_MoveDown[56] := BenchUut5.MoveDown;
   TraceOut_MoveUp[56] := BenchUut5.MoveUp;
   TraceOut_MoveLeft[56] := BenchUut5.MoveLeft;
   TraceOut_MoveRight[56] := BenchUut5.MoveRight;
   TraceOut_ActivateGrip[56] := BenchUut5.ActivateGrip;
   TraceOut_ActivateRelease[56] := BenchUut5.ActivateRelease;
   BenchCalls := BenchCalls + 1;
 57:
   BenchUut5.ManualMode := FALSE;
   BenchUut5.SingleStepMode := TRUE;
   BenchUut5.SingleCycleMode := FALSE;
   BenchUut5.ContinuousMode := FALSE;
   BenchUut5.EmergencyStop := TRUE;
   BenchUut5.Start := TRUE;
   BenchUut5.DownButton := FALSE;
   BenchUut5.UpButton := FALSE;
   BenchUut5.LeftButton := FALSE;
   BenchUut5.RightButton := FALSE;
   BenchUut5.GripButton := FALSE;
   BenchUut5.ReleaseButton := FALSE;
   BenchUut5.DownLimitSwitch := FALSE;
   BenchUut5.UpLimitSwitch := FALSE;
   BenchUut5.LeftLimitSwitch := FALSE;
   BenchUut5.RightLimitSwitch := FALSE;
   BenchUut5.GripLimitSwitch := FALSE;
   BenchUut5.ReleaseLimitSwitch := FALSE;
   TraceIn_ManualMode[57] := BenchUut5.ManualMode;
   TraceIn_SingleStepMode[57] := BenchUut5.SingleStepMode;
   TraceIn_SingleCycleMode[57] := BenchUut5.SingleCycleMode;
   TraceIn_ContinuousMode[57] := BenchUut5.ContinuousMode;
   TraceIn_EmergencyStop[57] := BenchUut5.EmergencyStop;
   TraceIn_Start[57] := BenchUut5.Start;
   TraceIn_DownButton[57] := BenchUut5.DownButton;
   TraceIn_UpButton[57] := BenchUut5.UpButton;
   TraceIn_LeftButton[57] := BenchUut5.LeftButton;
   TraceIn_RightButton[57] := BenchUut5.RightButton;
   TraceIn_GripButton[57] := BenchUut5.GripButton;
   TraceIn_ReleaseButton[57] := BenchUut5.ReleaseButton;
   TraceIn_DownLimitSwitch[57] := BenchUut5.DownLimitSwitch;
   TraceIn_UpLimitSwitch[57] := BenchUut5.UpLimitSwitch;
   TraceIn_LeftLimitSwitch[57] := BenchUut5.LeftLimitSwitch;
   TraceIn_RightLimitSwitch[57] := BenchUut5.RightLimitSwitch;
   TraceIn_GripLimitSwitch[57] := BenchUut5.GripLimitSwitch;
   TraceIn_ReleaseLimitSwitch[57] := BenchUut5.ReleaseLimitSwitch;
   BenchUut5();
   TraceOut_MoveDown[57] := BenchUut5.MoveDown;
   TraceOut_MoveUp[57] := BenchUut5.MoveUp;
   TraceOut_MoveLeft[57] := BenchUut5.MoveLeft;
   TraceOut_MoveRight[57] := BenchUut5.MoveRight;
   TraceOut_ActivateGrip[57] := BenchUut5.ActivateGrip;
   TraceOut_ActivateRelease[57] := BenchUut5.ActivateRelease;
   BenchCalls := BenchCalls + 1;
 58:
   BenchUut5.ManualMode := FALSE;
   BenchUut5.SingleStepMode := TRUE;
   BenchUut5.SingleCycleMode := FALSE;
   BenchUut5.ContinuousMode := FALSE;
   BenchUut5.EmergencyStop := TRUE;
   BenchUut5.Start := FALSE;
   BenchUut5.DownButton := FALSE;
   BenchUut5.UpButton := FALSE;
   BenchUut5.LeftButton := FALSE;
   BenchUut5.RightButton := FALSE;
   BenchUut5.GripButton := FALSE;
   BenchUut5.ReleaseButton := FALSE;
   BenchUut5.DownLimitSwitch := FALSE;
   BenchUut5.UpLimitSwitch := FALSE;
   BenchUut5.LeftLimitSwitch := FALSE;
   BenchUut5.RightLimitSwitch := TRUE;
   BenchUut5.GripLimitSwitch := FALSE;
   BenchUut5.ReleaseLimitSwitch := FALSE;
   TraceIn_ManualMode[58] := BenchUut5.ManualMode;
   TraceIn_SingleStepMode[58] := BenchUut5.SingleStepMode;
   TraceIn_SingleCycleMode[58] := BenchUut5.SingleCycleMode;
   TraceIn_ContinuousMode[58] := BenchUut5.ContinuousMode;
   TraceIn_EmergencyStop[58] := BenchUut5.EmergencyStop;
   TraceIn_Start[58] := BenchUut5.Start;
   TraceIn_DownButton[58] := BenchUut5.DownButton;
   TraceIn_UpButton[58] := BenchUut5.UpButton;
   TraceIn_LeftButton[58] := BenchUut5.LeftButton;
   TraceIn_RightButton[58] := BenchUut5.RightButton;
   TraceIn_GripButton[58] := BenchUut5.GripButton;
   TraceIn_ReleaseButton[58] := BenchUut5.ReleaseButton;
   TraceIn_DownLimitSwitch[58] := BenchUut5.DownLimitSwitch;
   TraceIn_UpLimitSwitch[58] := BenchUut5.UpLimitSwitch;
   TraceIn_LeftLimitSwitch[58] := BenchUut5.LeftLimitSwitch;
   TraceIn_RightLimitSwitch[58] := BenchUut5.RightLimitSwitch;
   TraceIn_GripLimitSwitch[58] := BenchUut5.GripLimitSwitch;
   TraceIn_ReleaseLimitSwitch[58] := BenchUut5.ReleaseLimitSwitch;
   BenchUut5();
   TraceOut_MoveDown[58] := BenchUut5.MoveDown;
   TraceOut_MoveUp[58] := BenchUut5.MoveUp;
   TraceOut_MoveLeft[58] := BenchUut5.MoveLeft;
   TraceOut_MoveRight[58] := BenchUut5.MoveRight;
   TraceOut_ActivateGrip[58] := BenchUut5.ActivateGrip;
   TraceOut_ActivateRelease[58] := BenchUut5.ActivateRelease;
   BenchCalls := BenchCalls + 1;
 59:
   BenchUut5.ManualMode := FALSE;
   BenchUut5.SingleStepMode := TRUE;
   BenchUut5.SingleCycleMode := FALSE;
   BenchUut5.ContinuousMode := FALSE;
   BenchUut5.EmergencyStop := TRUE;
   BenchUut5.Start := TRUE;
   BenchUut5.DownButton := FALSE;
   BenchUut5.UpButton := FALSE;
   BenchUut5.LeftButton := FALSE;
   BenchUut5.RightButton := FALSE;
   BenchUut5.GripButton := FALSE;
   BenchUut5.ReleaseButton := FALSE;
   BenchUut5.DownLimitSwitch := FALSE;
   BenchUut5.UpLimitSwitch := FALSE;
   BenchUut5.LeftLimitSwitch := FALSE;
   BenchUut5.RightLimitSwitch := FALSE;
   BenchUut5.GripLimitSwitch := FALSE;
   BenchUut5.ReleaseLimitSwitch := FALSE;
   TraceIn_ManualMode[59] := BenchUut5.ManualMode;
   TraceIn_SingleStepMode[59] := BenchUut5.SingleStepMode;
   TraceIn_SingleCycleMode[59] := BenchUut5.SingleCycleMode;
   TraceIn_ContinuousMode[59] := BenchUut5.ContinuousMode;
   TraceIn_EmergencyStop[59] := BenchUut5.EmergencyStop;
   TraceIn_Start[59] := BenchUut5.Start;
   TraceIn_DownButton[59] := BenchUut5.DownButton;
   TraceIn_UpButton[59] := BenchUut5.UpButton;
   TraceIn_LeftButton[59] := BenchUut5.LeftButton;
   TraceIn_RightButton[59] := BenchUut5.RightButton;
   TraceIn_GripButton[59] := BenchUut5.GripButton;
   TraceIn_ReleaseButton[59] := BenchUut5.ReleaseButton;
   TraceIn_DownLimitSwitch[59] := BenchUut5.DownLimitSwitch;
   TraceIn_UpLimitSwitch[59] := BenchUut5.UpLimitSwitch;
   TraceIn_LeftLimitSwitch[59] := BenchUut5.LeftLimitSwitch;
   TraceIn_RightLimitSwitch[59] := BenchUut5.RightLimitSwitch;
   TraceIn_GripLimitSwitch[59] := BenchUut5.GripLimitSwitch;
   TraceIn_ReleaseLimitSwitch[59] := BenchUut5.ReleaseLimitSwitch;
   BenchUut5();
   TraceOut_MoveDown[59] := BenchUut5.MoveDown;
   TraceOut_MoveUp[59] := BenchUut5.MoveUp;
   TraceOut_MoveLeft[59] := BenchUut5.MoveLeft;
   TraceOut_MoveRight[59] := BenchUut5.MoveRight;
   TraceOut_ActivateGrip[59] := BenchUut5.ActivateGrip;
   TraceOut_ActivateRelease[59] := BenchUut5.ActivateRelease;
   BenchCalls := BenchCalls + 1;
 60:
   BenchUut5.ManualMode := FALSE;
   BenchUut5.SingleStepMode := TRUE;
   BenchUut5.SingleCycleMode := FALSE;
   BenchUut5.ContinuousMode := FALSE;
   BenchUut5.EmergencyStop := TRUE;
   BenchUut5.Start := FALSE;
   BenchUut5.DownButton := FALSE;
   BenchUut5.UpButton := FALSE;
   BenchUut5.LeftButton := FALSE;
   BenchUut5.RightButton := FALSE;
   BenchUut5.GripButton := FALSE;
   BenchUut5.ReleaseButton := FALSE;
   BenchUut5.DownLimitSwitch := TRUE;
   BenchUut5.UpLimitSwitch := FALSE;
   BenchUut5.LeftLimitSwitch := FALSE;
   BenchUut5.RightLimitSwitch := FALSE;
   BenchUut5.GripLimitSwitch := FALSE;
   BenchUut5.ReleaseLimitSwitch := FALSE;
   TraceIn_ManualMode[60] := BenchUut5.ManualMode;
   TraceIn_SingleStepMode[60] := BenchUut5.SingleStepMode;
   TraceIn_SingleCycleMode[60] := BenchUut5.SingleCycleMode;
   TraceIn_ContinuousMode[60] := BenchUut5.ContinuousMode;
   TraceIn_EmergencyStop[60] := BenchUut5.EmergencyStop;
   TraceIn_Start[60] := BenchUut5.Start;
   TraceIn_DownButton[60] := BenchUut5.DownButton;
   TraceIn_UpButton[60] := BenchUut5.UpButton;
   TraceIn_LeftButton[60] := BenchUut5.LeftButton;
   TraceIn_RightButton[60] := BenchUut5.RightButton;
   TraceIn_GripButton[60] := BenchUut5.GripButton;
   TraceIn_ReleaseButton[60] := BenchUut5.ReleaseButton;
   TraceIn_DownLimitSwitch[60] := BenchUut5.DownLimitSwitch;
   TraceIn_UpLimitSwitch[60] := BenchUut5.UpLimitSwitch;
   TraceIn_LeftLimitSwitch[60] := BenchUut5.LeftLimitSwitch;
   TraceIn_RightLimitSwitch[60] := BenchUut5.RightLimitSwitch;
   TraceIn_GripLimitSwitch[60] := BenchUut5.GripLimitSwitch;
   TraceIn_ReleaseLimitSwitch[60] := BenchUut5.ReleaseLimitSwitch;
   BenchUut5();
   TraceOut_MoveDown[60] := BenchUut5.MoveDown;
   TraceOut_MoveUp[60] := BenchUut5.MoveUp;
   TraceOut_MoveLeft[60] := BenchUut5.MoveLeft;
   TraceOut_MoveRight[60] := BenchUut5.MoveRight;
   TraceOut_ActivateGrip[60] := BenchUut5.ActivateGrip;
   TraceOut_ActivateRelease[60] := BenchUut5.ActivateRelease;
   BenchCalls := BenchCalls + 1;
 61:
   BenchUut5.ManualMode := FALSE;
   BenchUut5.SingleStepMode := TRUE;
   BenchUut5.SingleCycleMode := FALSE;
   BenchUut5.ContinuousMode := FALSE;
   BenchUut5.EmergencyStop := TRUE;
   BenchUut5.Start := TRUE;
   BenchUut5.DownButton := FALSE;
   BenchUut5.UpButton := FALSE;
   BenchUut5.LeftButton := FALSE;
   BenchUut5.RightButton := FALSE;
   BenchUut5.GripButton := FALSE;
   BenchUut5.ReleaseButton := FALSE;
   BenchUut5.DownLimitSwitch := FALSE;
   BenchUut5.UpLimitSwitch := FALSE;
   BenchUut5.LeftLimitSwitch := FALSE;
   BenchUut5.RightLimitSwitch := FALSE;
   BenchUut5.GripLimitSwitch := FALSE;
   BenchUut5.ReleaseLimitSwitch := FALSE;
   TraceIn_ManualMode[61] := BenchUut5.ManualMode;
   TraceIn_SingleStepMode[61] := BenchUut5.SingleStepMode;
   TraceIn_SingleCycleMode[61] := BenchUut5.SingleCycleMode;
   TraceIn_ContinuousMode[61] := BenchUut5.ContinuousMode;
   TraceIn_EmergencyStop[61] := BenchUut5.EmergencyStop;
   TraceIn_Start[61] := BenchUut5.Start;
   TraceIn_DownButton[61] := BenchUut5.DownButton;
   TraceIn_UpButton[61] := BenchUut5.UpButton;
   TraceIn_LeftButton[61] := BenchUut5.LeftButton;
   TraceIn_RightButton[61] := BenchUut5.RightButton;
   TraceIn_GripButton[61] := BenchUut5.GripButton;
   TraceIn_ReleaseButton[61] := BenchUut5.ReleaseButton;
   TraceIn_DownLimitSwitch[61] := BenchUut5.DownLimitSwitch;
   TraceIn_UpLimitSwitch[61] := BenchUut5.UpLimitSwitch;
   TraceIn_LeftLimitSwitch[61] := BenchUut5.LeftLimitSwitch;
   TraceIn_RightLimitSwitch[61] := BenchUut5.RightLimitSwitch;
   TraceIn_GripLimitSwitch[61] := BenchUut5.GripLimitSwitch;
   TraceIn_ReleaseLimitSwitch[61] := BenchUut5.ReleaseLimitSwitch;
   BenchUut5();
   TraceOut_MoveDown[61] := BenchUut5.MoveDown;
   TraceOut_MoveUp[61] := BenchUut5.MoveUp;
   TraceOut_MoveLeft[61] := BenchUut5.MoveLeft;
   TraceOut_MoveRight[61] := BenchUut5.MoveRight;
   TraceOut_ActivateGrip[61] := BenchUut5.ActivateGrip;
   TraceOut_ActivateRelease[61] := BenchUut5.ActivateRelease;
   BenchCalls := BenchCalls + 1;
 62:
   BenchUut5.ManualMode := FALSE;
   BenchUut5.SingleStepMode := TRUE;
   BenchUut5.SingleCycleMode := FALSE;
   BenchUut5.ContinuousMode := FALSE;
   BenchUut5.EmergencyStop := TRUE;
   BenchUut5.Start := FALSE;
   BenchUut5.DownButton := FALSE;
   BenchUut5.UpButton := FALSE;
   BenchUut5.LeftButton := FALSE;
   BenchUut5.RightButton := FALSE;
   BenchUut5.GripButton := FALSE;
   BenchUut5.ReleaseButton := FALSE;
   BenchUut5.DownLimitSwitch := FALSE;
   BenchUut5.UpLimitSwitch := FALSE;
   BenchUut5.LeftLimitSwitch := FALSE;
   BenchUut5.RightLimitSwitch := FALSE;
   BenchUut5.GripLimitSwitch := FALSE;
   BenchUut5.ReleaseLimitSwitch := TRUE;
   TraceIn_ManualMode[62] := BenchUut5.ManualMode;
   TraceIn_SingleStepMode[62] := BenchUut5.SingleStepMode;
   TraceIn_SingleCycleMode[62] := BenchUut5.SingleCycleMode;
   TraceIn_ContinuousMode[62] := BenchUut5.ContinuousMode;
   TraceIn_EmergencyStop[62] := BenchUut5.EmergencyStop;
   TraceIn_Start[62] := BenchUut5.Start;
   TraceIn_DownButton[62] := BenchUut5.DownButton;
   TraceIn_UpButton[62] := BenchUut5.UpButton;
   TraceIn_LeftButton[62] := BenchUut5.LeftButton;
   TraceIn_RightButton[62] := BenchUut5.RightButton;
   TraceIn_GripButton[62] := BenchUut5.GripButton;
   TraceIn_ReleaseButton[62] := BenchUut5.ReleaseButton;
   TraceIn_DownLimitSwitch[62] := BenchUut5.DownLimitSwitch;
   TraceIn_UpLimitSwitch[62] := BenchUut5.UpLimitSwitch;
   TraceIn_LeftLimitSwitch[62] := BenchUut5.LeftLimitSwitch;
   TraceIn_RightLimitSwitch[62] := BenchUut5.RightLimitSwitch;
   TraceIn_GripLimitSwitch[62] := BenchUut5.GripLimitSwitch;
   TraceIn_ReleaseLimitSwitch[62] := BenchUut5.ReleaseLimitSwitch;
   BenchUut5();
   TraceOut_MoveDown[62] := BenchUut5.MoveDown;
   TraceOut_MoveUp[62] := BenchUut5.MoveUp;
   TraceOut_MoveLeft[62] := BenchUut5.MoveLeft;
   TraceOut_MoveRight[62] := BenchUut5.MoveRight;
   TraceOut_ActivateGrip[62] := BenchUut5.ActivateGrip;
   TraceOut_ActivateRelease[62] := BenchUut5.ActivateRelease;
   BenchCalls := BenchCalls + 1;
 63:
   BenchUut5.ManualMode := FALSE;
   BenchUut5.SingleStepMode := TRUE;
   BenchUut5.SingleCycleMode := FALSE;
   BenchUut5.ContinuousMode := FALSE;
   BenchUut5.EmergencyStop := TRUE;
   BenchUut5.Start := TRUE;
   BenchUut5.DownButton := FALSE;
   BenchUut5.UpButton := FALSE;
   BenchUut5.LeftButton := FALSE;
   BenchUut5.RightButton := FALSE;
   BenchUut5.GripButton := FALSE;
   BenchUut5.ReleaseButton := FALSE;
   BenchUut5.DownLimitSwitch := FALSE;
   BenchUut5.UpLimitSwitch := FALSE;
   BenchUut5.LeftLimitSwitch := FALSE;
   BenchUut5.RightLimitSwitch := FALSE;
   BenchUut5.GripLimitSwitch := FALSE;
   BenchUut5.ReleaseLimitSwitch := FALSE;
   TraceIn_ManualMode[63] := BenchUut5.ManualMode;
   TraceIn_SingleStepMode[63] := BenchUut5.SingleStepMode;
   TraceIn_SingleCycleMode[63] := BenchUut5.SingleCycleMode;
   TraceIn_ContinuousMode[63] := BenchUut5.ContinuousMode;
   TraceIn_EmergencyStop[63] := BenchUut5.EmergencyStop;
   TraceIn_Start[63] := BenchUut5.Start;
   TraceIn_DownButton[63] := BenchUut5.DownButton;
   TraceIn_UpButton[63] := BenchUut5.UpButton;
   TraceIn_LeftButton[63] := BenchUut5.LeftButton;
   TraceIn_RightButton[63] := BenchUut5.RightButton;
   TraceIn_GripButton[63] := BenchUut5.GripButton;
   TraceIn_ReleaseButton[63] := BenchUut5.ReleaseButton;
   TraceIn_DownLimitSwitch[63] := BenchUut5.DownLimitSwitch;
   TraceIn_UpLimitSwitch[63] := BenchUut5.UpLimitSwitch;
   TraceIn_LeftLimitSwitch[63] := BenchUut5.LeftLimitSwitch;
   TraceIn_RightLimitSwitch[63] := BenchUut5.RightLimitSwitch;
   TraceIn_GripLimitSwitch[63] := BenchUut5.GripLimitSwitch;
   TraceIn_ReleaseLimitSwitch[63] := BenchUut5.ReleaseLimitSwitch;
   BenchUut5();
   TraceOut_MoveDown[63] := BenchUut5.MoveDown;
   TraceOut_MoveUp[63] := BenchUut5.MoveUp;
   TraceOut_MoveLeft[63] := BenchUut5.MoveLeft;
   TraceOut_MoveRight[63] := BenchUut5.MoveRight;
   TraceOut_ActivateGrip[63] := BenchUut5.ActivateGrip;
   TraceOut_ActivateRelease[63] := BenchUut5.ActivateRelease;
   BenchCalls := BenchCalls + 1;
 64:
   BenchUut5.ManualMode := FALSE;
   BenchUut5.SingleStepMode := TRUE;
   BenchUut5.SingleCycleMode := FALSE;
   BenchUut5.ContinuousMode := FALSE;
   BenchUut5.EmergencyStop := TRUE;
   BenchUut5.Start := FALSE;
   BenchUut5.DownButton := FALSE;
   BenchUut5.UpButton := FALSE;
   BenchUut5.LeftButton := FALSE;
   BenchUut5.RightButton := FALSE;
   BenchUut5.GripButton := FALSE;
   BenchUut5.ReleaseButton := FALSE;
   BenchUut5.DownLimitSwitch := FALSE;
   BenchUut5.UpLimitSwitch := TRUE;
   BenchUut5.LeftLimitSwitch := FALSE;
   BenchUut5.RightLimitSwitch := FALSE;
   BenchUut5.GripLimitSwitch := FALSE;
   BenchUut5.ReleaseLimitSwitch := FALSE;
   TraceIn_ManualMode[64] := BenchUut5.ManualMode;
   TraceIn_SingleStepMode[64] := BenchUut5.SingleStepMode;
   TraceIn_SingleCycleMode[64] := BenchUut5.SingleCycleMode;
   TraceIn_ContinuousMode[64] := BenchUut5.ContinuousMode;
   TraceIn_EmergencyStop[64] := BenchUut5.EmergencyStop;
   TraceIn_Start[64] := BenchUut5.Start;
   TraceIn_DownButton[64] := BenchUut5.DownButton;
   TraceIn_UpButton[64] := BenchUut5.UpButton;
   TraceIn_LeftButton[64] := BenchUut5.LeftButton;
   TraceIn_RightButton[64] := BenchUut5.RightButton;
   TraceIn_GripButton[64] := BenchUut5.GripButton;
   TraceIn_ReleaseButton[64] := BenchUut5.ReleaseButton;
   TraceIn_DownLimitSwitch[64] := BenchUut5.DownLimitSwitch;
   TraceIn_UpLimitSwitch[64] := BenchUut5.UpLimitSwitch;
   TraceIn_LeftLimitSwitch[64] := BenchUut5.LeftLimitSwitch;
   TraceIn_RightLimitSwitch[64] := BenchUut5.RightLimitSwitch;
   TraceIn_GripLimitSwitch[64] := BenchUut5.GripLimitSwitch;
   TraceIn_ReleaseLimitSwitch[64] := BenchUut5.ReleaseLimitSwitch;
   BenchUut5();
   TraceOut_MoveDown[64] := BenchUut5.MoveDown;
   TraceOut_MoveUp[64] := BenchUut5.MoveUp;
   TraceOut_MoveLeft[64] := BenchUut5.MoveLeft;
   TraceOut_MoveRight[64] := BenchUut5.MoveRight;
   TraceOut_ActivateGrip[64] := BenchUut5.ActivateGrip;
   TraceOut_ActivateRelease[64] := BenchUut5.ActivateRelease;
   BenchCalls := BenchCalls + 1;
 65:
   BenchUut5.ManualMode := FALSE;
   BenchUut5.SingleStepMode := TRUE;
   BenchUut5.SingleCycleMode := FALSE;
   BenchUut5.ContinuousMode := FALSE;
   BenchUut5.EmergencyStop := TRUE;
   BenchUut5.Start := TRUE;
   BenchUut5.DownButton := FALSE;
   BenchUut5.UpButton := FALSE;
   BenchUut5.LeftButton := FALSE;
   BenchUut5.RightButton := FALSE;
   BenchUut5.GripButton := FALSE;
   BenchUut5.ReleaseButton := FALSE;
   BenchUut5.DownLimitSwitch := FALSE;
   BenchUut5.UpLimitSwitch := FALSE;
   BenchUut5.LeftLimitSwitch := FALSE;
   BenchUut5.RightLimitSwitch := FALSE;
   BenchUut5.GripLimitSwitch := FALSE;
   BenchUut5.ReleaseLimitSwitch := FALSE;
   TraceIn_ManualMode[65] := BenchUut5.ManualMode;
   TraceIn_SingleStepMode[65] := BenchUut5.SingleStepMode;
   TraceIn_SingleCycleMode[65] := BenchUut5.SingleCycleMode;
   TraceIn_ContinuousMode[65] := BenchUut5.ContinuousMode;
   TraceIn_EmergencyStop[65] := BenchUut5.EmergencyStop;
   TraceIn_Start[65] := BenchUut5.Start;
   TraceIn_DownButton[65] := BenchUut5.DownButton;
   TraceIn_UpButton[65] := BenchUut5.UpButton;
   TraceIn_LeftButton[65] := BenchUut5.LeftButton;
   TraceIn_RightButton[65] := BenchUut5.RightButton;
   TraceIn_GripButton[65] := BenchUut5.GripButton;
   TraceIn_ReleaseButton[65] := BenchUut5.ReleaseButton;
   TraceIn_DownLimitSwitch[65] := BenchUut5.DownLimitSwitch;
   TraceIn_UpLimitSwitch[65] := BenchUut5.UpLimitSwitch;
   TraceIn_LeftLimitSwitch[65] := BenchUut5.LeftLimitSwitch;
   TraceIn_RightLimitSwitch[65] := BenchUut5.RightLimitSwitch;
   TraceIn_GripLimitSwitch[65] := BenchUut5.GripLimitSwitch;
   TraceIn_ReleaseLimitSwitch[65] := BenchUut5.ReleaseLimitSwitch;
   BenchUut5();
   TraceOut_MoveDown[65] := BenchUut5.MoveDown;
   TraceOut_MoveUp[65] := BenchUut5.MoveUp;
   TraceOut_MoveLeft[65] := BenchUut5.MoveLeft;
   TraceOut_MoveRight[65] := BenchUut5.MoveRight;
   TraceOut_ActivateGrip[65] := BenchUut5.ActivateGrip;
   TraceOut_ActivateRelease[65] := BenchUut5.ActivateRelease;
   BenchCalls := BenchCalls + 1;
 66:
   BenchUut5.ManualMode := FALSE;
   BenchUut5.SingleStepMode := TRUE;
   BenchUut5.SingleCycleMode := FALSE;
   BenchUut5.ContinuousMode := FALSE;
   BenchUut5.EmergencyStop := TRUE;
   BenchUut5.Start := FALSE;
   BenchUut5.DownButton := FALSE;
   BenchUut5.UpButton := FALSE;
   BenchUut5.LeftButton := FALSE;
   BenchUut5.RightButton := FALSE;
   BenchUut5.GripButton := FALSE;
   BenchUut5.ReleaseButton := FALSE;
   BenchUut5.DownLimitSwitch := FALSE;
   BenchUut5.UpLimitSwitch := TRUE;
   BenchUut5.LeftLimitSwitch := TRUE;
   BenchUut5.RightLimitSwitch := FALSE;
   BenchUut5.GripLimitSwitch := FALSE;
   BenchUut5.ReleaseLimitSwitch := FALSE;
   TraceIn_ManualMode[66] := BenchUut5.ManualMode;
   TraceIn_SingleStepMode[66] := BenchUut5.SingleStepMode;
   TraceIn_SingleCycleMode[66] := BenchUut5.SingleCycleMode;
   TraceIn_ContinuousMode[66] := BenchUut5.ContinuousMode;
   TraceIn_EmergencyStop[66] := BenchUut5.EmergencyStop;
   TraceIn_Start[66] := BenchUut5.Start;
   TraceIn_DownButton[66] := BenchUut5.DownButton;
   TraceIn_UpButton[66] := BenchUut5.UpButton;
   TraceIn_LeftButton[66] := BenchUut5.LeftButton;
   TraceIn_RightButton[66] := BenchUut5.RightButton;
   TraceIn_GripButton[66] := BenchUut5.GripButton;
   TraceIn_ReleaseButton[66] := BenchUut5.ReleaseButton;
   TraceIn_DownLimitSwitch[66] := BenchUut5.DownLimitSwitch;
   TraceIn_UpLimitSwitch[66] := BenchUut5.UpLimitSwitch;
   TraceIn_LeftLimitSwitch[66] := BenchUut5.LeftLimitSwitch;
   TraceIn_RightLimitSwitch[66] := BenchUut5.RightLimitSwitch;
   TraceIn_GripLimitSwitch[66] := BenchUut5.GripLimitSwitch;
   TraceIn_ReleaseLimitSwitch[66] := BenchUut5.ReleaseLimitSwitch;
   BenchUut5();
   TraceOut_MoveDown[66] := BenchUut5.MoveDown;
   TraceOut_MoveUp[66] := BenchUut5.MoveUp;
   TraceOut_MoveLeft[66] := BenchUut5.MoveLeft;
   TraceOut_MoveRight[66] := BenchUut5.MoveRight;
   TraceOut_ActivateGrip[66] := BenchUut5.ActivateGrip;
   TraceOut_ActivateRelease[66] := BenchUut5.ActivateRelease;
   BenchCalls := BenchCalls + 1;
 67:
   BenchUut5.ManualMode := FALSE;
   BenchUut5.SingleStepMode := TRUE;
   BenchUut5.SingleCycleMode := FALSE;
   BenchUut5.ContinuousMode := FALSE;
   BenchUut5.EmergencyStop := FALSE;
   BenchUut5.Start := FALSE;
   BenchUut5.DownButton := FALSE;
   BenchUut5.UpButton := FALSE;
   BenchUut5.LeftButton := FALSE;
   BenchUut5.RightButton := FALSE;
   BenchUut5.GripButton := FALSE;
   BenchUut5.ReleaseButton := FALSE;
   BenchUut5.DownLimitSwitch := FALSE;
   BenchUut5.UpLimitSwitch := FALSE;
   BenchUut5.LeftLimitSwitch := FALSE;
   BenchUut5.RightLimitSwitch := FALSE;
   BenchUut5.GripLimitSwitch := FALSE;
   BenchUut5.ReleaseLimitSwitch := FALSE;
   TraceIn_ManualMode[67] := BenchUut5.ManualMode;
   TraceIn_SingleStepMode[67] := BenchUut5.SingleStepMode;
   TraceIn_SingleCycleMode[67] := BenchUut5.SingleCycleMode;
   TraceIn_ContinuousMode[67] := BenchUut5.ContinuousMode;
   TraceIn_EmergencyStop[67] := BenchUut5.EmergencyStop;
   TraceIn_Start[67] := BenchUut5.Start;
   TraceIn_DownButton[67] := BenchUut5.DownButton;
   TraceIn_UpButton[67] := BenchUut5.UpButton;
   TraceIn_LeftButton[67] := BenchUut5.LeftButton;
   TraceIn_RightButton[67] := BenchUut5.RightButton;
   TraceIn_GripButton[67] := BenchUut5.GripButton;
   TraceIn_ReleaseButton[67] := BenchUut5.ReleaseButton;
   TraceIn_DownLimitSwitch[67] := BenchUut5.DownLimitSwitch;
   TraceIn_UpLimitSwitch[67] := BenchUut5.UpLimitSwitch;
   TraceIn_LeftLimitSwitch[67] := BenchUut5.LeftLimitSwitch;
   TraceIn_RightLimitSwitch[67] := BenchUut5.RightLimitSwitch;
   TraceIn_GripLimitSwitch[67] := BenchUut5.GripLimitSwitch;
   TraceIn_ReleaseLimitSwitch[67] := BenchUut5.ReleaseLimitSwitch;
   BenchUut5();
   TraceOut_MoveDown[67] := BenchUut5.MoveDown;
   TraceOut_MoveUp[67] := BenchUut5.MoveUp;
   TraceOut_MoveLeft[67] := BenchUut5.MoveLeft;
   TraceOut_MoveRight[67] := BenchUut5.MoveRight;
   TraceOut_ActivateGrip[67] := BenchUut5.ActivateGrip;
   TraceOut_ActivateRelease[67] := BenchUut5.ActivateRelease;
   BenchCalls := BenchCalls + 1;
 68:
   BenchUut5.ManualMode := TRUE;
   BenchUut5.SingleStepMode := FALSE;
   BenchUut5.SingleCycleMode := FALSE;
   BenchUut5.ContinuousMode := FALSE;
   BenchUut5.EmergencyStop := TRUE;
   BenchUut5.Start := FALSE;
   BenchUut5.DownButton := FALSE;
   BenchUut5.UpButton := FALSE;
   BenchUut5.LeftButton := FALSE;
   BenchUut5.RightButton := TRUE;
   BenchUut5.GripButton := FALSE;
   BenchUut5.ReleaseButton := FALSE;
   BenchUut5.DownLimitSwitch := FALSE;
   BenchUut5.UpLimitSwitch := FALSE;
   BenchUut5.LeftLimitSwitch := FALSE;
   BenchUut5.RightLimitSwitch := FALSE;
   BenchUut5.GripLimitSwitch := FALSE;
   BenchUut5.ReleaseLimitSwitch := FALSE;
   TraceIn_ManualMode[68] := BenchUut5.ManualMode;
   TraceIn_SingleStepMode[68] := BenchUut5.SingleStepMode;
   TraceIn_SingleCycleMode[68] := BenchUut5.SingleCycleMode;
   TraceIn_ContinuousMode[68] := BenchUut5.ContinuousMode;
   TraceIn_EmergencyStop[68] := BenchUut5.EmergencyStop;
   TraceIn_Start[68] := BenchUut5.Start;
   TraceIn_DownButton[68] := BenchUut5.DownButton;
   TraceIn_UpButton[68] := BenchUut5.UpButton;
   TraceIn_LeftButton[68] := BenchUut5.LeftButton;
   TraceIn_RightButton[68] := BenchUut5.RightButton;
   TraceIn_GripButton[68] := BenchUut5.GripButton;
   TraceIn_ReleaseButton[68] := BenchUut5.ReleaseButton;
   TraceIn_DownLimitSwitch[68] := BenchUut5.DownLimitSwitch;
   TraceIn_UpLimitSwitch[68] := BenchUut5.UpLimitSwitch;
   TraceIn_LeftLimitSwitch[68] := BenchUut5.LeftLimitSwitch;
   TraceIn_RightLimitSwitch[68] := BenchUut5.RightLimitSwitch;
   TraceIn_GripLimitSwitch[68] := BenchUut5.GripLimitSwitch;
   TraceIn_ReleaseLimitSwitch[68] := BenchUut5.ReleaseLimitSwitch;
   BenchUut5();
   TraceOut_MoveDown[68] := BenchUut5.MoveDown;
   TraceOut_MoveUp[68] := BenchUut5.MoveUp;
   TraceOut_MoveLeft[68] := BenchUut5.MoveLeft;
   TraceOut_MoveRight[68] := BenchUut5.MoveRight;
   TraceOut_ActivateGrip[68] := BenchUut5.ActivateGrip;
   TraceOut_ActivateRelease[68] := BenchUut5.ActivateRelease;
   BenchCalls := BenchCalls + 1;
 69:
   BenchUut5.ManualMode := TRUE;
   BenchUut5.SingleStepMode := FALSE;
   BenchUut5.SingleCycleMode := FALSE;
   BenchUut5.ContinuousMode := FALSE;
   BenchUut5.EmergencyStop := TRUE;
   BenchUut5.Start := FALSE;
   BenchUut5.DownButton := FALSE;
   BenchUut5.UpButton := FALSE;
   BenchUut5.LeftButton := FALSE;
   BenchUut5.RightButton := TRUE;
   BenchUut5.GripButton := FALSE;
   BenchUut5.ReleaseButton := FALSE;
   BenchUut5.DownLimitSwitch := FALSE;
   BenchUut5.UpLimitSwitch := FALSE;
   BenchUut5.LeftLimitSwitch := FALSE;
   BenchUut5.RightLimitSwitch := FALSE;
   BenchUut5.GripLimitSwitch := FALSE;
   BenchUut5.ReleaseLimitSwitch := FALSE;
   TraceIn_ManualMode[69] := BenchUut5.ManualMode;
   TraceIn_SingleStepMode[69] := BenchUut5.SingleStepMode;
   TraceIn_SingleCycleMode[69] := BenchUut5.SingleCycleMode;
   TraceIn_ContinuousMode[69] := BenchUut5.ContinuousMode;
   TraceIn_EmergencyStop[69] := BenchUut5.EmergencyStop;
   TraceIn_Start[69] := BenchUut5.Start;
   TraceIn_DownButton[69] := BenchUut5.DownButton;
   TraceIn_UpButton[69] := BenchUut5.UpButton;
   TraceIn_LeftButton[69] := BenchUut5.LeftButton;
   TraceIn_RightButton[69] := BenchUut5.RightButton;
   TraceIn_GripButton[69] := BenchUut5.GripButton;
   TraceIn_ReleaseButton[69] := BenchUut5.ReleaseButton;
   TraceIn_DownLimitSwitch[69] := BenchUut5.DownLimitSwitch;
   TraceIn_UpLimitSwitch[69] := BenchUut5.UpLimitSwitch;
   TraceIn_LeftLimitSwitch[69] := BenchUut5.LeftLimitSwitch;
   TraceIn_RightLimitSwitch[69] := BenchUut5.RightLimitSwitch;
   TraceIn_GripLimitSwitch[69] := BenchUut5.GripLimitSwitch;
   TraceIn_ReleaseLimitSwitch[69] := BenchUut5.ReleaseLimitSwitch;
   BenchUut5();
   TraceOut_MoveDown[69] := BenchUut5.MoveDown;
   TraceOut_MoveUp[69] := BenchUut5.MoveUp;
   TraceOut_MoveLeft[69] := BenchUut5.MoveLeft;
   TraceOut_MoveRight[69] := BenchUut5.MoveRight;
   TraceOut_ActivateGrip[69] := BenchUut5.ActivateGrip;
   TraceOut_ActivateRelease[69] := BenchUut5.ActivateRelease;
   BenchCalls := BenchCalls + 1;
 70:
   BenchUut6.ManualMode := TRUE;
   BenchUut6.SingleStepMode := FALSE;
   BenchUut6.SingleCycleMode := FALSE;
   BenchUut6.ContinuousMode := FALSE;
   BenchUut6.EmergencyStop := TRUE;
   BenchUut6.Start := FALSE;
   BenchUut6.DownButton := FALSE;
   BenchUut6.UpButton := TRUE;
   BenchUut6.LeftButton := FALSE;
   BenchUut6.RightButton := FALSE;
   BenchUut6.GripButton := FALSE;
   BenchUut6.ReleaseButton := FALSE;
   BenchUut6.DownLimitSwitch := FALSE;
   BenchUut6.UpLimitSwitch := FALSE;
   BenchUut6.LeftLimitSwitch := TRUE;
   BenchUut6.RightLimitSwitch := FALSE;
   BenchUut6.GripLimitSwitch := FALSE;
   BenchUut6.ReleaseLimitSwitch := TRUE;
   TraceIn_ManualMode[70] := BenchUut6.ManualMode;
   TraceIn_SingleStepMode[70] := BenchUut6.SingleStepMode;
   TraceIn_SingleCycleMode[70] := BenchUut6.SingleCycleMode;
   TraceIn_ContinuousMode[70] := BenchUut6.ContinuousMode;
   TraceIn_EmergencyStop[70] := BenchUut6.EmergencyStop;
   TraceIn_Start[70] := BenchUut6.Start;
   TraceIn_DownButton[70] := BenchUut6.DownButton;
   TraceIn_UpButton[70] := BenchUut6.UpButton;
   TraceIn_LeftButton[70] := BenchUut6.LeftButton;
   TraceIn_RightButton[70] := BenchUut6.RightButton;
   TraceIn_GripButton[70] := BenchUut6.GripButton;
   TraceIn_ReleaseButton[70] := BenchUut6.ReleaseButton;
   TraceIn_DownLimitSwitch[70] := BenchUut6.DownLimitSwitch;
   TraceIn_UpLimitSwitch[70] := BenchUut6.UpLimitSwitch;
   TraceIn_LeftLimitSwitch[70] := BenchUut6.LeftLimitSwitch;
   TraceIn_RightLimitSwitch[70] := BenchUut6.RightLimitSwitch;
   TraceIn_GripLimitSwitch[70] := BenchUut6.GripLimitSwitch;
   TraceIn_ReleaseLimitSwitch[70] := BenchUut6.ReleaseLimitSwitch;
   BenchUut6();
   TraceOut_MoveDown[70] := BenchUut6.MoveDown;
   TraceOut_MoveUp[70] := BenchUut6.MoveUp;
   TraceOut_MoveLeft[70] := BenchUut6.MoveLeft;
   TraceOut_MoveRight[70] := BenchUut6.MoveRight;
   TraceOut_ActivateGrip[70] := BenchUut6.ActivateGrip;
   TraceOut_ActivateRelease[70] := BenchUut6.ActivateRelease;
   BenchCalls := BenchCalls + 1;
 71:
   BenchUut7.ManualMode := FALSE;
   BenchUut7.SingleStepMode := FALSE;
   BenchUut7.SingleCycleMode := TRUE;
   BenchUut7.ContinuousMode := FALSE;
   BenchUut7.EmergencyStop := TRUE;
   BenchUut7.Start := FALSE;
   BenchUut7.DownButton := FALSE;
   BenchUut7.UpButton := FALSE;
   BenchUut7.LeftButton := FALSE;
   BenchUut7.RightButton := FALSE;
   BenchUut7.GripButton := FALSE;
   BenchUut7.ReleaseButton := FALSE;
   BenchUut7.DownLimitSwitch := FALSE;
   BenchUut7.UpLimitSwitch := TRUE;
   BenchUut7.LeftLimitSwitch := TRUE;
   BenchUut7.RightLimitSwitch := FALSE;
   BenchUut7.GripLimitSwitch := FALSE;
   BenchUut7.ReleaseLimitSwitch := TRUE;
   TraceIn_ManualMode[71] := BenchUut7.ManualMode;
   TraceIn_SingleStepMode[71] := BenchUut7.SingleStepMode;
   TraceIn_SingleCycleMode[71] := BenchUut7.SingleCycleMode;
   TraceIn_ContinuousMode[71] := BenchUut7.ContinuousMode;
   TraceIn_EmergencyStop[71] := BenchUut7.EmergencyStop;
   TraceIn_Start[71] := BenchUut7.Start;
   TraceIn_DownButton[71] := BenchUut7.DownButton;
   TraceIn_UpButton[71] := BenchUut7.UpButton;
   TraceIn_LeftButton[71] := BenchUut7.LeftButton;
   TraceIn_RightButton[71] := BenchUut7.RightButton;
   TraceIn_GripButton[71] := BenchUut7.GripButton;
   TraceIn_ReleaseButton[71] := BenchUut7.ReleaseButton;
   TraceIn_DownLimitSwitch[71] := BenchUut7.DownLimitSwitch;
   TraceIn_UpLimitSwitch[71] := BenchUut7.UpLimitSwitch;
   TraceIn_LeftLimitSwitch[71] := BenchUut7.LeftLimitSwitch;
   TraceIn_RightLimitSwitch[71] := BenchUut7.RightLimitSwitch;
   TraceIn_GripLimitSwitch[71] := BenchUut7.GripLimitSwitch;
   TraceIn_ReleaseLimitSwitch[71] := BenchUut7.ReleaseLimitSwitch;
   BenchUut7();
   TraceOut_MoveDown[71] := BenchUut7.MoveDown;
   TraceOut_MoveUp[71] := BenchUut7.MoveUp;
   TraceOut_MoveLeft[71] := BenchUut7.MoveLeft;
   TraceOut_MoveRight[71] := BenchUut7.MoveRight;
   TraceOut_ActivateGrip[71] := BenchUut7.ActivateGrip;
   TraceOut_ActivateRelease[71] := BenchUut7.ActivateRelease;
   BenchCalls := BenchCalls + 1;
 72:
   BenchUut7.ManualMode := FALSE;
   BenchUut7.SingleStepMode := FALSE;
   BenchUut7.SingleCycleMode := TRUE;
   BenchUut7.ContinuousMode := FALSE;
   BenchUut7.EmergencyStop := TRUE;
   BenchUut7.Start := TRUE;
   BenchUut7.DownButton := FALSE;
   BenchUut7.UpButton := FALSE;
   BenchUut7.LeftButton := FALSE;
   BenchUut7.RightButton := FALSE;
   BenchUut7.GripButton := FALSE;
   BenchUut7.ReleaseButton := FALSE;
   BenchUut7.DownLimitSwitch := FALSE;
   BenchUut7.UpLimitSwitch := TRUE;
   BenchUut7.LeftLimitSwitch := TRUE;
   BenchUut7.RightLimitSwitch := FALSE;
   BenchUut7.GripLimitSwitch := FALSE;
   BenchUut7.ReleaseLimitSwitch := TRUE;
   TraceIn_ManualMode[72] := BenchUut7.ManualMode;
   TraceIn_SingleStepMode[72] := BenchUut7.SingleStepMode;
   TraceIn_SingleCycleMode[72] := BenchUut7.SingleCycleMode;
   TraceIn_ContinuousMode[72] := BenchUut7.ContinuousMode;
   TraceIn_EmergencyStop[72] := BenchUut7.EmergencyStop;
   TraceIn_Start[72] := BenchUut7.Start;
   TraceIn_DownButton[72] := BenchUut7.DownButton;
   TraceIn_UpButton[72] := BenchUut7.UpButton;
   TraceIn_LeftButton[72] := BenchUut7.LeftButton;
   TraceIn_RightButton[72] := BenchUut7.RightButton;
   TraceIn_GripButton[72] := BenchUut7.GripButton;
   TraceIn_ReleaseButton[72] := BenchUut7.ReleaseButton;
   TraceIn_DownLimitSwitch[72] := BenchUut7.DownLimitSwitch;
   TraceIn_UpLimitSwitch[72] := BenchUut7.UpLimitSwitch;
   TraceIn_LeftLimitSwitch[72] := BenchUut7.LeftLimitSwitch;
   TraceIn_RightLimitSwitch[72] := BenchUut7.RightLimitSwitch;
   TraceIn_GripLimitSwitch[72] := BenchUut7.GripLimitSwitch;
   TraceIn_ReleaseLimitSwitch[72] := BenchUut7.ReleaseLimitSwitch;
   BenchUut7();
   TraceOut_MoveDown[72] := BenchUut7.MoveDown;
   TraceOut_MoveUp[72] := BenchUut7.MoveUp;
   TraceOut_MoveLeft[72] := BenchUut7.MoveLeft;
   TraceOut_MoveRight[72] := BenchUut7.MoveRight;
   TraceOut_ActivateGrip[72] := BenchUut7.ActivateGrip;
   TraceOut_ActivateRelease[72] := BenchUut7.ActivateRelease;
   BenchCalls := BenchCalls + 1;
 73:
   BenchUut7.ManualMode := FALSE;
   BenchUut7.SingleStepMode := FALSE;
   BenchUut7.SingleCycleMode := TRUE;
   BenchUut7.ContinuousMode := FALSE;
   BenchUut7.EmergencyStop := TRUE;
   BenchUut7.Start := FALSE;
   BenchUut7.DownButton := FALSE;
   BenchUut7.UpButton := FALSE;
   BenchUut7.LeftButton := FALSE;
   BenchUut7.RightButton := FALSE;
   BenchUut7.GripButton := FALSE;
   BenchUut7.ReleaseButton := FALSE;
   BenchUut7.DownLimitSwitch := TRUE;
   BenchUut7.UpLimitSwitch := FALSE;
   BenchUut7.LeftLimitSwitch := TRUE;
   BenchUut7.RightLimitSwitch := FALSE;
   BenchUut7.GripLimitSwitch := FALSE;
   BenchUut7.ReleaseLimitSwitch := FALSE;
   TraceIn_ManualMode[73] := BenchUut7.ManualMode;
   TraceIn_SingleStepMode[73] := BenchUut7.SingleStepMode;
   TraceIn_SingleCycleMode[73] := BenchUut7.SingleCycleMode;
   TraceIn_ContinuousMode[73] := BenchUut7.ContinuousMode;
   TraceIn_EmergencyStop[73] := BenchUut7.EmergencyStop;
   TraceIn_Start[73] := BenchUut7.Start;
   TraceIn_DownButton[73] := BenchUut7.DownButton;
   TraceIn_UpButton[73] := BenchUut7.UpButton;
   TraceIn_LeftButton[73] := BenchUut7.LeftButton;
   TraceIn_RightButton[73] := BenchUut7.RightButton;
   TraceIn_GripButton[73] := BenchUut7.GripButton;
   TraceIn_ReleaseButton[73] := BenchUut7.ReleaseButton;
   TraceIn_DownLimitSwitch[73] := BenchUut7.DownLimitSwitch;
   TraceIn_UpLimitSwitch[73] := BenchUut7.UpLimitSwitch;
   TraceIn_LeftLimitSwitch[73] := BenchUut7.LeftLimitSwitch;
   TraceIn_RightLimitSwitch[73] := BenchUut7.RightLimitSwitch;
   TraceIn_GripLimitSwitch[73] := BenchUut7.GripLimitSwitch;
   TraceIn_ReleaseLimitSwitch[73] := BenchUut7.ReleaseLimitSwitch;
   BenchUut7();
   TraceOut_MoveDown[73] := BenchUut7.MoveDown;
   TraceOut_MoveUp[73] := BenchUut7.MoveUp;
   TraceOut_MoveLeft[73] := BenchUut7.MoveLeft;
   TraceOut_MoveRight[73] := BenchUut7.MoveRight;
   TraceOut_ActivateGrip[73] := BenchUut7.ActivateGrip;
   TraceOut_ActivateRelease[73] := BenchUut7.ActivateRelease;
   BenchCalls := BenchCalls + 1;
 74:
   BenchUut7.ManualMode := FALSE;
   BenchUut7.SingleStepMode := FALSE;
   BenchUut7.SingleCycleMode := TRUE;
   BenchUut7.ContinuousMode := FALSE;
   BenchUut7.EmergencyStop := TRUE;
   BenchUut7.Start := FALSE;
   BenchUut7.DownButton := FALSE;
   BenchUut7.UpButton := FALSE;
   BenchUut7.LeftButton := FALSE;
   BenchUut7.RightButton := FALSE;
   BenchUut7.GripButton := FALSE;
   BenchUut7.ReleaseButton := FALSE;
   BenchUut7.DownLimitSwitch := TRUE;
   BenchUut7.UpLimitSwitch := FALSE;
   BenchUut7.LeftLimitSwitch := TRUE;
   BenchUut7.RightLimitSwitch := FALSE;
   BenchUut7.GripLimitSwitch := FALSE;
   BenchUut7.ReleaseLimitSwitch := FALSE;
   TraceIn_ManualMode[74] := BenchUut7.ManualMode;
   TraceIn_SingleStepMode[74] := BenchUut7.SingleStepMode;
   TraceIn_SingleCycleMode[74] := BenchUut7.SingleCycleMode;
   TraceIn_ContinuousMode[74] := BenchUut7.ContinuousMode;
   TraceIn_EmergencyStop[74] := BenchUut7.EmergencyStop;
   TraceIn_Start[74] := BenchUut7.Start;
   TraceIn_DownButton[74] := BenchUut7.DownButton;
   TraceIn_UpButton[74] := BenchUut7.UpButton;
   TraceIn_LeftButton[74] := BenchUut7.LeftButton;
   TraceIn_RightButton[74] := BenchUut7.RightButton;
   TraceIn_GripButton[74] := BenchUut7.GripButton;
   TraceIn_ReleaseButton[74] := BenchUut7.ReleaseButton;
   TraceIn_DownLimitSwitch[74] := BenchUut7.DownLimitSwitch;
   TraceIn_UpLimitSwitch[74] := BenchUut7.UpLimitSwitch;
   TraceIn_LeftLimitSwitch[74] := BenchUut7.LeftLimitSwitch;
   TraceIn_RightLimitSwitch[74] := BenchUut7.RightLimitSwitch;
   TraceIn_GripLimitSwitch[74] := BenchUut7.GripLimitSwitch;
   TraceIn_ReleaseLimitSwitch[74] := BenchUut7.ReleaseLimitSwitch;
   BenchUut7();
   TraceOut_MoveDown[74] := BenchUut7.MoveDown;
   TraceOut_MoveUp[74] := BenchUut7.MoveUp;
   TraceOut_MoveLeft[74] := BenchUut7.MoveLeft;
   TraceOut_MoveRight[74] := BenchUut7.MoveRight;
   TraceOut_ActivateGrip[74] := BenchUut7.ActivateGrip;
   TraceOut_ActivateRelease[74] := BenchUut7.ActivateRelease;
   BenchCalls := BenchCalls + 1;
 75:
   BenchUut8.ManualMode := TRUE;
   BenchUut8.SingleStepMode := FALSE;
   BenchUut8.SingleCycleMode := FALSE;
   BenchUut8.ContinuousMode := FALSE;
   BenchUut8.EmergencyStop := TRUE;
   BenchUut8.Start := FALSE;
   BenchUut8.DownButton := FALSE;
   BenchUut8.UpButton := FALSE;
   BenchUut8.LeftButton := FALSE;
   BenchUut8.RightButton := FALSE;
   BenchUut8.GripButton := FALSE;
   BenchUut8.ReleaseButton := FALSE;
   BenchUut8.DownLimitSwitch := FALSE;
   BenchUut8.UpLimitSwitch := FALSE;
   BenchUut8.LeftLimitSwitch := FALSE;
   BenchUut8.RightLimitSwitch := FALSE;
   BenchUut8.GripLimitSwitch := FALSE;
   BenchUut8.ReleaseLimitSwitch := FALSE;
   TraceIn_ManualMode[75] := BenchUut8.ManualMode;
   TraceIn_SingleStepMode[75] := BenchUut8.SingleStepMode;
   TraceIn_SingleCycleMode[75] := BenchUut8.SingleCycleMode;
   TraceIn_ContinuousMode[75] := BenchUut8.ContinuousMode;
   TraceIn_EmergencyStop[75] := BenchUut8.EmergencyStop;
   TraceIn_Start[75] := BenchUut8.Start;
   TraceIn_DownButton[75] := BenchUut8.DownButton;
   TraceIn_UpButton[75] := BenchUut8.UpButton;
   TraceIn_LeftButton[75] := BenchUut8.LeftButton;
   TraceIn_RightButton[75] := BenchUut8.RightButton;
   TraceIn_GripButton[75] := BenchUut8.GripButton;
   TraceIn_ReleaseButton[75] := BenchUut8.ReleaseButton;
   TraceIn_DownLimitSwitch[75] := BenchUut8.DownLimitSwitch;
   TraceIn_UpLimitSwitch[75] := BenchUut8.UpLimitSwitch;
   TraceIn_LeftLimitSwitch[75] := BenchUut8.LeftLimitSwitch;
   TraceIn_RightLimitSwitch[75] := BenchUut8.RightLimitSwitch;
   TraceIn_GripLimitSwitch[75] := BenchUut8.GripLimitSwitch;
   TraceIn_ReleaseLimitSwitch[75] := BenchUut8.ReleaseLimitSwitch;
   BenchUut8();
   TraceOut_MoveDown[75] := BenchUut8.MoveDown;
   TraceOut_MoveUp[75] := BenchUut8.MoveUp;
   TraceOut_MoveLeft[75] := BenchUut8.MoveLeft;
   TraceOut_MoveRight[75] := BenchUut8.MoveRight;
   TraceOut_ActivateGrip[75] := BenchUut8.ActivateGrip;
   TraceOut_ActivateRelease[75] := BenchUut8.ActivateRelease;
   BenchCalls := BenchCalls + 1;
 76:
   BenchUut8.ManualMode := TRUE;
   BenchUut8.SingleStepMode := FALSE;
   BenchUut8.SingleCycleMode := FALSE;
   BenchUut8.ContinuousMode := FALSE;
   BenchUut8.EmergencyStop := TRUE;
   BenchUut8.Start := FALSE;
   BenchUut8.DownButton := TRUE;
   BenchUut8.UpButton := FALSE;
   BenchUut8.LeftButton := FALSE;
   BenchUut8.RightButton := FALSE;
   BenchUut8.GripButton := FALSE;
   BenchUut8.ReleaseButton := FALSE;
   BenchUut8.DownLimitSwitch := FALSE;
   BenchUut8.UpLimitSwitch := FALSE;
   BenchUut8.LeftLimitSwitch := FALSE;
   BenchUut8.RightLimitSwitch := FALSE;
   BenchUut8.GripLimitSwitch := FALSE;
   BenchUut8.ReleaseLimitSwitch := FALSE;
   TraceIn_ManualMode[76] := BenchUut8.ManualMode;
   TraceIn_SingleStepMode[76] := BenchUut8.SingleStepMode;
   TraceIn_SingleCycleMode[76] := BenchUut8.SingleCycleMode;
   TraceIn_ContinuousMode[76] := BenchUut8.ContinuousMode;
   TraceIn_EmergencyStop[76] := BenchUut8.EmergencyStop;
   TraceIn_Start[76] := BenchUut8.Start;
   TraceIn_DownButton[76] := BenchUut8.DownButton;
   TraceIn_UpButton[76] := BenchUut8.UpButton;
   TraceIn_LeftButton[76] := BenchUut8.LeftButton;
   TraceIn_RightButton[76] := BenchUut8.RightButton;
   TraceIn_GripButton[76] := BenchUut8.GripButton;
   TraceIn_ReleaseButton[76] := BenchUut8.ReleaseButton;
   TraceIn_DownLimitSwitch[76] := BenchUut8.DownLimitSwitch;
   TraceIn_UpLimitSwitch[76] := BenchUut8.UpLimitSwitch;
   TraceIn_LeftLimitSwitch[76] := BenchUut8.LeftLimitSwitch;
   TraceIn_RightLimitSwitch[76] := BenchUut8.RightLimitSwitch;
   TraceIn_GripLimitSwitch[76] := BenchUut8.GripLimitSwitch;
   TraceIn_ReleaseLimitSwitch[76] := BenchUut8.ReleaseLimitSwitch;
   BenchUut8();
   TraceOut_MoveDown[76] := BenchUut8.MoveDown;
   TraceOut_MoveUp[76] := BenchUut8.MoveUp;
   TraceOut_MoveLeft[76] := BenchUut8.MoveLeft;
   TraceOut_MoveRight[76] := BenchUut8.MoveRight;
   TraceOut_ActivateGrip[76] := BenchUut8.ActivateGrip;
   TraceOut_ActivateRelease[76] := BenchUut8.ActivateRelease;
   BenchCalls := BenchCalls + 1;
 77:
   BenchUut8.ManualMode := TRUE;
   BenchUut8.SingleStepMode := FALSE;
   BenchUut8.SingleCycleMode := FALSE;
   BenchUut8.ContinuousMode := FALSE;
   BenchUut8.EmergencyStop := TRUE;
   BenchUut8.Start := FALSE;
   BenchUut8.DownButton := TRUE;
   BenchUut8.UpButton := FALSE;
   BenchUut8.LeftButton := FALSE;
   BenchUut8.RightButton := FALSE;
   BenchUut8.GripButton := FALSE;
   BenchUut8.ReleaseButton := FALSE;
   BenchUut8.DownLimitSwitch := FALSE;
   BenchUut8.UpLimitSwitch := FALSE;
   BenchUut8.LeftLimitSwitch := FALSE;
   BenchUut8.RightLimitSwitch := FALSE;
   BenchUut8.GripLimitSwitch := FALSE;
   BenchUut8.ReleaseLimitSwitch := FALSE;
   TraceIn_ManualMode[77] := BenchUut8.ManualMode;
   TraceIn_SingleStepMode[77] := BenchUut8.SingleStepMode;
   TraceIn_SingleCycleMode[77] := BenchUut8.SingleCycleMode;
   TraceIn_ContinuousMode[77] := BenchUut8.ContinuousMode;
   TraceIn_EmergencyStop[77] := BenchUut8.EmergencyStop;
   TraceIn_Start[77] := BenchUut8.Start;
   TraceIn_DownButton[77] := BenchUut8.DownButton;
   TraceIn_UpButton[77] := BenchUut8.UpButton;
   TraceIn_LeftButton[77] := BenchUut8.LeftButton;
   TraceIn_RightButton[77] := BenchUut8.RightButton;
   TraceIn_GripButton[77] := BenchUut8.GripButton;
   TraceIn_ReleaseButton[77] := BenchUut8.ReleaseButton;
   TraceIn_DownLimitSwitch[77] := BenchUut8.DownLimitSwitch;
   TraceIn_UpLimitSwitch[77] := BenchUut8.UpLimitSwitch;
   TraceIn_LeftLimitSwitch[77] := BenchUut8.LeftLimitSwitch;
   TraceIn_RightLimitSwitch[77] := BenchUut8.RightLimitSwitch;
   TraceIn_GripLimitSwitch[77] := BenchUut8.GripLimitSwitch;
   TraceIn_ReleaseLimitSwitch[77] := BenchUut8.ReleaseLimitSwitch;
   BenchUut8();
   TraceOut_MoveDown[77] := BenchUut8.MoveDown;
   TraceOut_MoveUp[77] := BenchUut8.MoveUp;
   TraceOut_MoveLeft[77] := BenchUut8.MoveLeft;
   TraceOut_MoveRight[77] := BenchUut8.MoveRight;
   TraceOut_ActivateGrip[77] := BenchUut8.ActivateGrip;
   TraceOut_ActivateRelease[77] := BenchUut8.ActivateRelease;
   BenchCalls := BenchCalls + 1;
 78:
   BenchUut8.ManualMode := TRUE;
   BenchUut8.SingleStepMode := FALSE;
   BenchUut8.SingleCycleMode := FALSE;
   BenchUut8.ContinuousMode := FALSE;
   BenchUut8.EmergencyStop := TRUE;
   BenchUut8.Start := FALSE;
   BenchUut8.DownButton := TRUE;
   BenchUut8.UpButton := FALSE;
   BenchUut8.LeftButton := FALSE;
   BenchUut8.RightButton := FALSE;
   BenchUut8.GripButton := FALSE;
   BenchUut8.ReleaseButton := FALSE;
   BenchUut8.DownLimitSwitch := TRUE;
   BenchUut8.UpLimitSwitch := FALSE;
   BenchUut8.LeftLimitSwitch := FALSE;
   BenchUut8.RightLimitSwitch := FALSE;
   BenchUut8.GripLimitSwitch := FALSE;
   BenchUut8.ReleaseLimitSwitch := FALSE;
   TraceIn_ManualMode[78] := BenchUut8.ManualMode;
   TraceIn_SingleStepMode[78] := BenchUut8.SingleStepMode;
   TraceIn_SingleCycleMode[78] := BenchUut8.SingleCycleMode;
   TraceIn_ContinuousMode[78] := BenchUut8.ContinuousMode;
   TraceIn_EmergencyStop[78] := BenchUut8.EmergencyStop;
   TraceIn_Start[78] := BenchUut8.Start;
   TraceIn_DownButton[78] := BenchUut8.DownButton;
   TraceIn_UpButton[78] := BenchUut8.UpButton;
   TraceIn_LeftButton[78] := BenchUut8.LeftButton;
   TraceIn_RightButton[78] := BenchUut8.RightButton;
   TraceIn_GripButton[78] := BenchUut8.GripButton;
   TraceIn_ReleaseButton[78] := BenchUut8.ReleaseButton;
   TraceIn_DownLimitSwitch[78] := BenchUut8.DownLimitSwitch;
   TraceIn_UpLimitSwitch[78] := BenchUut8.UpLimitSwitch;
   TraceIn_LeftLimitSwitch[78] := BenchUut8.LeftLimitSwitch;
   TraceIn_RightLimitSwitch[78] := BenchUut8.RightLimitSwitch;
   TraceIn_GripLimitSwitch[78] := BenchUut8.GripLimitSwitch;
   TraceIn_ReleaseLimitSwitch[78] := BenchUut8.ReleaseLimitSwitch;
   BenchUut8();
   TraceOut_MoveDown[78] := BenchUut8.MoveDown;
   TraceOut_MoveUp[78] := BenchUut8.MoveUp;
   TraceOut_MoveLeft[78] := BenchUut8.MoveLeft;
   TraceOut_MoveRight[78] := BenchUut8.MoveRight;
   TraceOut_ActivateGrip[78] := BenchUut8.ActivateGrip;
   TraceOut_ActivateRelease[78] := BenchUut8.ActivateRelease;
   BenchCalls := BenchCalls + 1;
 79:
   BenchUut8.ManualMode := TRUE;
   BenchUut8.SingleStepMode := FALSE;
   BenchUut8.SingleCycleMode := FALSE;
   BenchUut8.ContinuousMode := FALSE;
   BenchUut8.EmergencyStop := TRUE;
   BenchUut8.Start := FALSE;
   BenchUut8.DownButton := FALSE;
   BenchUut8.UpButton := FALSE;
   BenchUut8.LeftButton := FALSE;
   BenchUut8.RightButton := FALSE;
   BenchUut8.GripButton := FALSE;
   BenchUut8.ReleaseButton := FALSE;
   BenchUut8.DownLimitSwitch := TRUE;
   BenchUut8.UpLimitSwitch := FALSE;
   BenchUut8.LeftLimitSwitch := FALSE;
   BenchUut8.RightLimitSwitch := FALSE;
   BenchUut8.GripLimitSwitch := FALSE;
   BenchUut8.ReleaseLimitSwitch := FALSE;
   TraceIn_ManualMode[79] := BenchUut8.ManualMode;
   TraceIn_SingleStepMode[79] := BenchUut8.SingleStepMode;
   TraceIn_SingleCycleMode[79] := BenchUut8.SingleCycleMode;
   TraceIn_ContinuousMode[79] := BenchUut8.ContinuousMode;
   TraceIn_EmergencyStop[79] := BenchUut8.EmergencyStop;
   TraceIn_Start[79] := BenchUut8.Start;
   TraceIn_DownButton[79] := BenchUut8.DownButton;
   TraceIn_UpButton[79] := BenchUut8.UpButton;
   TraceIn_LeftButton[79] := BenchUut8.LeftButton;
   TraceIn_RightButton[79] := BenchUut8.RightButton;
   TraceIn_GripButton[79] := BenchUut8.GripButton;
   TraceIn_ReleaseButton[79] := BenchUut8.ReleaseButton;
   TraceIn_DownLimitSwitch[79] := BenchUut8.DownLimitSwitch;
   TraceIn_UpLimitSwitch[79] := BenchUut8.UpLimitSwitch;
   TraceIn_LeftLimitSwitch[79] := BenchUut8.LeftLimitSwitch;
   TraceIn_RightLimitSwitch[79] := BenchUut8.RightLimitSwitch;
   TraceIn_GripLimitSwitch[79] := BenchUut8.GripLimitSwitch;
   TraceIn_ReleaseLimitSwitch[79] := BenchUut8.ReleaseLimitSwitch;
   BenchUut8();
   TraceOut_MoveDown[79] := BenchUut8.MoveDown;
   TraceOut_MoveUp[79] := BenchUut8.MoveUp;
   TraceOut_MoveLeft[79] := BenchUut8.MoveLeft;
   TraceOut_MoveRight[79] := BenchUut8.MoveRight;
   TraceOut_ActivateGrip[79] := BenchUut8.ActivateGrip;
   TraceOut_ActivateRelease[79] := BenchUut8.ActivateRelease;
   BenchCalls := BenchCalls + 1;
 80:
   BenchUut8.ManualMode := TRUE;
   BenchUut8.SingleStepMode := FALSE;
   BenchUut8.SingleCycleMode := FALSE;
   BenchUut8.ContinuousMode := FALSE;
   BenchUut8.EmergencyStop := TRUE;
   BenchUut8.Start := FALSE;
   BenchUut8.DownButton := FALSE;
   BenchUut8.UpButton := FALSE;
   BenchUut8.LeftButton := FALSE;
   BenchUut8.RightButton := FALSE;
   BenchUut8.GripButton := FALSE;
   BenchUut8.ReleaseButton := FALSE;
   BenchUut8.DownLimitSwitch := FALSE;
   BenchUut8.UpLimitSwitch := FALSE;
   BenchUut8.LeftLimitSwitch := FALSE;
   BenchUut8.RightLimitSwitch := FALSE;
   BenchUut8.GripLimitSwitch := FALSE;
   BenchUut8.ReleaseLimitSwitch := FALSE;
   TraceIn_ManualMode[80] := BenchUut8.ManualMode;
   TraceIn_SingleStepMode[80] := BenchUut8.SingleStepMode;
   TraceIn_SingleCycleMode[80] := BenchUut8.SingleCycleMode;
   TraceIn_ContinuousMode[80] := BenchUut8.ContinuousMode;
   TraceIn_EmergencyStop[80] := BenchUut8.EmergencyStop;
   TraceIn_Start[80] := BenchUut8.Start;
   TraceIn_DownButton[80] := BenchUut8.DownButton;
   TraceIn_UpButton[80] := BenchUut8.UpButton;
   TraceIn_LeftButton[80] := BenchUut8.LeftButton;
   TraceIn_RightButton[80] := BenchUut8.RightButton;
   TraceIn_GripButton[80] := BenchUut8.GripButton;
   TraceIn_ReleaseButton[80] := BenchUut8.ReleaseButton;
   TraceIn_DownLimitSwitch[80] := BenchUut8.DownLimitSwitch;
   TraceIn_UpLimitSwitch[80] := BenchUut8.UpLimitSwitch;
   TraceIn_LeftLimitSwitch[80] := BenchUut8.LeftLimitSwitch;
   TraceIn_RightLimitSwitch[80] := BenchUut8.RightLimitSwitch;
   TraceIn_GripLimitSwitch[80] := BenchUut8.GripLimitSwitch;
   TraceIn_ReleaseLimitSwitch[80] := BenchUut8.ReleaseLimitSwitch;
   BenchUut8();
   TraceOut_MoveDown[80] := BenchUut8.MoveDown;
   TraceOut_MoveUp[80] := BenchUut8.MoveUp;
   TraceOut_MoveLeft[80] := BenchUut8.MoveLeft;
   TraceOut_MoveRight[80] := BenchUut8.MoveRight;
   TraceOut_ActivateGrip[80] := BenchUut8.ActivateGrip;
   TraceOut_ActivateRelease[80] := BenchUut8.ActivateRelease;
   BenchCalls := BenchCalls + 1;
 81:
   BenchUut9.ManualMode := TRUE;
   BenchUut9.SingleStepMode := FALSE;
   BenchUut9.SingleCycleMode := FALSE;
   BenchUut9.ContinuousMode := FALSE;
   BenchUut9.EmergencyStop := TRUE;
   BenchUut9.Start := FALSE;
   BenchUut9.DownButton := FALSE;
   BenchUut9.UpButton := FALSE;
   BenchUut9.LeftButton := FALSE;
   BenchUut9.RightButton := FALSE;
   BenchUut9.GripButton := FALSE;
   BenchUut9.ReleaseButton := FALSE;
   BenchUut9.DownLimitSwitch := FALSE;
   BenchUut9.UpLimitSwitch := FALSE;
   BenchUut9.LeftLimitSwitch := FALSE;
   BenchUut9.RightLimitSwitch := FALSE;
   BenchUut9.GripLimitSwitch := FALSE;
   BenchUut9.ReleaseLimitSwitch := FALSE;
   TraceIn_ManualMode[81] := BenchUut9.ManualMode;
   TraceIn_SingleStepMode[81] := BenchUut9.SingleStepMode;
   TraceIn_SingleCycleMode[81] := BenchUut9.SingleCycleMode;
   TraceIn_ContinuousMode[81] := BenchUut9.ContinuousMode;
   TraceIn_EmergencyStop[81] := BenchUut9.EmergencyStop;
   TraceIn_Start[81] := BenchUut9.Start;
   TraceIn_DownButton[81] := BenchUut9.DownButton;
   TraceIn_UpButton[81] := BenchUut9.UpButton;
   TraceIn_LeftButton[81] := BenchUut9.LeftButton;
   TraceIn_RightButton[81] := BenchUut9.RightButton;
   TraceIn_GripButton[81] := BenchUut9.GripButton;
   TraceIn_ReleaseButton[81] := BenchUut9.ReleaseButton;
   TraceIn_DownLimitSwitch[81] := BenchUut9.DownLimitSwitch;
   TraceIn_UpLimitSwitch[81] := BenchUut9.UpLimitSwitch;
   TraceIn_LeftLimitSwitch[81] := BenchUut9.LeftLimitSwitch;
   TraceIn_RightLimitSwitch[81] := BenchUut9.RightLimitSwitch;
   TraceIn_GripLimitSwitch[81] := BenchUut9.GripLimitSwitch;
   TraceIn_ReleaseLimitSwitch[81] := BenchUut9.ReleaseLimitSwitch;
   BenchUut9();
   TraceOut_MoveDown[81] := BenchUut9.MoveDown;
   TraceOut_MoveUp[81] := BenchUut9.MoveUp;
   TraceOut_MoveLeft[81] := BenchUut9.MoveLeft;
   TraceOut_MoveRight[81] := BenchUut9.MoveRight;
   TraceOut_ActivateGrip[81] := BenchUut9.ActivateGrip;
   TraceOut_ActivateRelease[81] := BenchUut9.ActivateRelease;
   BenchCalls := BenchCalls + 1;
 82:
   BenchUut9.ManualMode := TRUE;
   BenchUut9.SingleStepMode := FALSE;
   BenchUut9.SingleCycleMode := FALSE;
   BenchUut9.ContinuousMode := FALSE;
   BenchUut9.EmergencyStop := TRUE;
   BenchUut9.Start := FALSE;
   BenchUut9.DownButton := FALSE;
   BenchUut9.UpButton := TRUE;
   BenchUut9.LeftButton := FALSE;
   BenchUut9.RightButton := FALSE;
   BenchUut9.GripButton := FALSE;
   BenchUut9.ReleaseButton := FALSE;
   BenchUut9.DownLimitSwitch := FALSE;
   BenchUut9.UpLimitSwitch := FALSE;
   BenchUut9.LeftLimitSwitch := FALSE;
   BenchUut9.RightLimitSwitch := FALSE;
   BenchUut9.GripLimitSwitch := FALSE;
   BenchUut9.ReleaseLimitSwitch := FALSE;
   TraceIn_ManualMode[82] := BenchUut9.ManualMode;
   TraceIn_SingleStepMode[82] := BenchUut9.SingleStepMode;
   TraceIn_SingleCycleMode[82] := BenchUut9.SingleCycleMode;
   TraceIn_ContinuousMode[82] := BenchUut9.ContinuousMode;
   TraceIn_EmergencyStop[82] := BenchUut9.EmergencyStop;
   TraceIn_Start[82] := BenchUut9.Start;
   TraceIn_DownButton[82] := BenchUut9.DownButton;
   TraceIn_UpButton[82] := BenchUut9.UpButton;
   TraceIn_LeftButton[82] := BenchUut9.LeftButton;
   TraceIn_RightButton[82] := BenchUut9.RightButton;
   TraceIn_GripButton[82] := BenchUut9.GripButton;
   TraceIn_ReleaseButton[82] := BenchUut9.ReleaseButton;
   TraceIn_DownLimitSwitch[82] := BenchUut9.DownLimitSwitch;
   TraceIn_UpLimitSwitch[82] := BenchUut9.UpLimitSwitch;
   TraceIn_LeftLimitSwitch[82] := BenchUut9.LeftLimitSwitch;
   TraceIn_RightLimitSwitch[82] := BenchUut9.RightLimitSwitch;
   TraceIn_GripLimitSwitch[82] := BenchUut9.GripLimitSwitch;
   TraceIn_ReleaseLimitSwitch[82] := BenchUut9.ReleaseLimitSwitch;
   BenchUut9();
   TraceOut_MoveDown[82] := BenchUut9.MoveDown;
   TraceOut_MoveUp[82] := BenchUut9.MoveUp;
   TraceOut_MoveLeft[82] := BenchUut9.MoveLeft;
   TraceOut_MoveRight[82] := BenchUut9.MoveRight;
   TraceOut_ActivateGrip[82] := BenchUut9.ActivateGrip;
   TraceOut_ActivateRelease[82] := BenchUut9.ActivateRelease;
   BenchCalls := BenchCalls + 1;
 83:
   BenchUut9.ManualMode := TRUE;
   BenchUut9.SingleStepMode := FALSE;
   BenchUut9.SingleCycleMode := FALSE;
   BenchUut9.ContinuousMode := FALSE;
   BenchUut9.EmergencyStop := TRUE;
   BenchUut9.Start := FALSE;
   BenchUut9.DownButton := FALSE;
   BenchUut9.UpButton := TRUE;
   BenchUut9.LeftButton := FALSE;
   BenchUut9.RightButton := FALSE;
   BenchUut9.GripButton := FALSE;
   BenchUut9.ReleaseButton := FALSE;
   BenchUut9.DownLimitSwitch := FALSE;
   BenchUut9.UpLimitSwitch := FALSE;
   BenchUut9.LeftLimitSwitch := FALSE;
   BenchUut9.RightLimitSwitch := FALSE;
   BenchUut9.GripLimitSwitch := FALSE;
   BenchUut9.ReleaseLimitSwitch := FALSE;
   TraceIn_ManualMode[83] := BenchUut9.ManualMode;
   TraceIn_SingleStepMode[83] := BenchUut9.SingleStepMode;
   TraceIn_SingleCycleMode[83] := BenchUut9.SingleCycleMode;
   TraceIn_ContinuousMode[83] := BenchUut9.ContinuousMode;
   TraceIn_EmergencyStop[83] := BenchUut9.EmergencyStop;
   TraceIn_Start[83] := BenchUut9.Start;
   TraceIn_DownButton[83] := BenchUut9.DownButton;
   TraceIn_UpButton[83] := BenchUut9.UpButton;
   TraceIn_LeftButton[83] := BenchUut9.LeftButton;
   TraceIn_RightButton[83] := BenchUut9.RightButton;
   TraceIn_GripButton[83] := BenchUut9.GripButton;
   TraceIn_ReleaseButton[83] := BenchUut9.ReleaseButton;
   TraceIn_DownLimitSwitch[83] := BenchUut9.DownLimitSwitch;
   TraceIn_UpLimitSwitch[83] := BenchUut9.UpLimitSwitch;
   TraceIn_LeftLimitSwitch[83] := BenchUut9.LeftLimitSwitch;
   TraceIn_RightLimitSwitch[83] := BenchUut9.RightLimitSwitch;
   TraceIn_GripLimitSwitch[83] := BenchUut9.GripLimitSwitch;
   TraceIn_ReleaseLimitSwitch[83] := BenchUut9.ReleaseLimitSwitch;
   BenchUut9();
   TraceOut_MoveDown[83] := BenchUut9.MoveDown;
   TraceOut_MoveUp[83] := BenchUut9.MoveUp;
   TraceOut_MoveLeft[83] := BenchUut9.MoveLeft;
   TraceOut_MoveRight[83] := BenchUut9.MoveRight;
   TraceOut_ActivateGrip[83] := BenchUut9.ActivateGrip;
   TraceOut_ActivateRelease[83] := BenchUut9.ActivateRelease;
   BenchCalls := BenchCalls + 1;
 84:
   BenchUut9.ManualMode := TRUE;
   BenchUut9.SingleStepMode := FALSE;
   BenchUut9.SingleCycleMode := FALSE;
   BenchUut9.ContinuousMode := FALSE;
   BenchUut9.EmergencyStop := TRUE;
   BenchUut9.Start := FALSE;
   BenchUut9.DownButton := FALSE;
   BenchUut9.UpButton := TRUE;
   BenchUut9.LeftButton := FALSE;
   BenchUut9.RightButton := FALSE;
   BenchUut9.GripButton := FALSE;
   BenchUut9.ReleaseButton := FALSE;
   BenchUut9.DownLimitSwitch := FALSE;
   BenchUut9.UpLimitSwitch := TRUE;
   BenchUut9.LeftLimitSwitch := FALSE;
   BenchUut9.RightLimitSwitch := FALSE;
   BenchUut9.GripLimitSwitch := FALSE;
   BenchUut9.ReleaseLimitSwitch := FALSE;
   TraceIn_ManualMode[84] := BenchUut9.ManualMode;
   TraceIn_SingleStepMode[84] := BenchUut9.SingleStepMode;
   TraceIn_SingleCycleMode[84] := BenchUut9.SingleCycleMode;
   TraceIn_ContinuousMode[84] := BenchUut9.ContinuousMode;
   TraceIn_EmergencyStop[84] := BenchUut9.EmergencyStop;
   TraceIn_Start[84] := BenchUut9.Start;
   TraceIn_DownButton[84] := BenchUut9.DownButton;
   TraceIn_UpButton[84] := BenchUut9.UpButton;
   TraceIn_LeftButton[84] := BenchUut9.LeftButton;
   TraceIn_RightButton[84] := BenchUut9.RightButton;
   TraceIn_GripButton[84] := BenchUut9.GripButton;
   TraceIn_ReleaseButton[84] := BenchUut9.ReleaseButton;
   TraceIn_DownLimitSwitch[84] := BenchUut9.DownLimitSwitch;
   TraceIn_UpLimitSwitch[84] := BenchUut9.UpLimitSwitch;
   TraceIn_LeftLimitSwitch[84] := BenchUut9.LeftLimitSwitch;
   TraceIn_RightLimitSwitch[84] := BenchUut9.RightLimitSwitch;
   TraceIn_GripLimitSwitch[84] := BenchUut9.GripLimitSwitch;
   TraceIn_ReleaseLimitSwitch[84] := BenchUut9.ReleaseLimitSwitch;
   BenchUut9();
   TraceOut_MoveDown[84] := BenchUut9.MoveDown;
   TraceOut_MoveUp[84] := BenchUut9.MoveUp;
   TraceOut_MoveLeft[84] := BenchUut9.MoveLeft;
   TraceOut_MoveRight[84] := BenchUut9.MoveRight;
   TraceOut_ActivateGrip[84] := BenchUut9.ActivateGrip;
   TraceOut_ActivateRelease[84] := BenchUut9.ActivateRelease;
   BenchCalls := BenchCalls + 1;
 85:
   BenchUut9.ManualMode := TRUE;
   BenchUut9.SingleStepMode := FALSE;
   BenchUut9.SingleCycleMode := FALSE;
   BenchUut9.ContinuousMode := FALSE;
   BenchUut9.EmergencyStop := TRUE;
   BenchUut9.Start := FALSE;
   BenchUut9.DownButton := FALSE;
   BenchUut9.UpButton := FALSE;
   BenchUut9.LeftButton := FALSE;
   BenchUut9.RightButton := FALSE;
   BenchUut9.GripButton := FALSE;
   BenchUut9.ReleaseButton := FALSE;
   BenchUut9.DownLimitSwitch := FALSE;
   BenchUut9.UpLimitSwitch := TRUE;
   BenchUut9.LeftLimitSwitch := FALSE;
   BenchUut9.RightLimitSwitch := FALSE;
   BenchUut9.GripLimitSwitch := FALSE;
   BenchUut9.ReleaseLimitSwitch := FALSE;
   TraceIn_ManualMode[85] := BenchUut9.ManualMode;
   TraceIn_SingleStepMode[85] := BenchUut9.SingleStepMode;
   TraceIn_SingleCycleMode[85] := BenchUut9.SingleCycleMode;
   TraceIn_ContinuousMode[85] := BenchUut9.ContinuousMode;
   TraceIn_EmergencyStop[85] := BenchUut9.EmergencyStop;
   TraceIn_Start[85] := BenchUut9.Start;
   TraceIn_DownButton[85] := BenchUut9.DownButton;
   TraceIn_UpButton[85] := BenchUut9.UpButton;
   TraceIn_LeftButton[85] := BenchUut9.LeftButton;
   TraceIn_RightButton[85] := BenchUut9.RightButton;
   TraceIn_GripButton[85] := BenchUut9.GripButton;
   TraceIn_ReleaseButton[85] := BenchUut9.ReleaseButton;
   TraceIn_DownLimitSwitch[85] := BenchUut9.DownLimitSwitch;
   TraceIn_UpLimitSwitch[85] := BenchUut9.UpLimitSwitch;
   TraceIn_LeftLimitSwitch[85] := BenchUut9.LeftLimitSwitch;
   TraceIn_RightLimitSwitch[85] := BenchUut9.RightLimitSwitch;
   TraceIn_GripLimitSwitch[85] := BenchUut9.GripLimitSwitch;
   TraceIn_ReleaseLimitSwitch[85] := BenchUut9.ReleaseLimitSwitch;
   BenchUut9();
   TraceOut_MoveDown[85] := BenchUut9.MoveDown;
   TraceOut_MoveUp[85] := BenchUut9.MoveUp;
   TraceOut_MoveLeft[85] := BenchUut9.MoveLeft;
   TraceOut_MoveRight[85] := BenchUut9.MoveRight;
   TraceOut_ActivateGrip[85] := BenchUut9.ActivateGrip;
   TraceOut_ActivateRelease[85] := BenchUut9.ActivateRelease;
   BenchCalls := BenchCalls + 1;
 86:
   BenchUut9.ManualMode := TRUE;
   BenchUut9.SingleStepMode := FALSE;
   BenchUut9.SingleCycleMode := FALSE;
   BenchUut9.ContinuousMode := FALSE;
   BenchUut9.EmergencyStop := TRUE;
   BenchUut9.Start := FALSE;
   BenchUut9.DownButton := FALSE;
   BenchUut9.UpButton := FALSE;
   BenchUut9.LeftButton := FALSE;
   BenchUut9.RightButton := FALSE;
   BenchUut9.GripButton := FALSE;
   BenchUut9.ReleaseButton := FALSE;
   BenchUut9.DownLimitSwitch := FALSE;
   BenchUut9.UpLimitSwitch := FALSE;
   BenchUut9.LeftLimitSwitch := FALSE;
   BenchUut9.RightLimitSwitch := FALSE;
   BenchUut9.GripLimitSwitch := FALSE;
   BenchUut9.ReleaseLimitSwitch := FALSE;
   TraceIn_ManualMode[86] := BenchUut9.ManualMode;
   TraceIn_SingleStepMode[86] := BenchUut9.SingleStepMode;
   TraceIn_SingleCycleMode[86] := BenchUut9.SingleCycleMode;
   TraceIn_ContinuousMode[86] := BenchUut9.ContinuousMode;
   TraceIn_EmergencyStop[86] := BenchUut9.EmergencyStop;
   TraceIn_Start[86] := BenchUut9.Start;
   TraceIn_DownButton[86] := BenchUut9.DownButton;
   TraceIn_UpButton[86] := BenchUut9.UpButton;
   TraceIn_LeftButton[86] := BenchUut9.LeftButton;
   TraceIn_RightButton[86] := BenchUut9.RightButton;
   TraceIn_GripButton[86] := BenchUut9.GripButton;
   TraceIn_ReleaseButton[86] := BenchUut9.ReleaseButton;
   TraceIn_DownLimitSwitch[86] := BenchUut9.DownLimitSwitch;
   TraceIn_UpLimitSwitch[86] := BenchUut9.UpLimitSwitch;
   TraceIn_LeftLimitSwitch[86] := BenchUut9.LeftLimitSwitch;
   TraceIn_RightLimitSwitch[86] := BenchUut9.RightLimitSwitch;
   TraceIn_GripLimitSwitch[86] := BenchUut9.GripLimitSwitch;
   TraceIn_ReleaseLimitSwitch[86] := BenchUut9.ReleaseLimitSwitch;
   BenchUut9();
   TraceOut_MoveDown[86] := BenchUut9.MoveDown;
   TraceOut_MoveUp[86] := BenchUut9.MoveUp;
   TraceOut_MoveLeft[86] := BenchUut9.MoveLeft;
   TraceOut_MoveRight[86] := BenchUut9.MoveRight;
   TraceOut_ActivateGrip[86] := BenchUut9.ActivateGrip;
   TraceOut_ActivateRelease[86] := BenchUut9.ActivateRelease;
   BenchCalls := BenchCalls + 1;
 87:
   BenchUut10.ManualMode := TRUE;
   BenchUut10.SingleStepMode := FALSE;
   BenchUut10.SingleCycleMode := FALSE;
   BenchUut10.ContinuousMode := FALSE;
   BenchUut10.EmergencyStop := TRUE;
   BenchUut10.Start := FALSE;
   BenchUut10.DownButton := FALSE;
   BenchUut10.UpButton := FALSE;
   BenchUut10.LeftButton := FALSE;
   BenchUut10.RightButton := FALSE;
   BenchUut10.GripButton := FALSE;
   BenchUut10.ReleaseButton := FALSE;
   BenchUut10.DownLimitSwitch := FALSE;
   BenchUut10.UpLimitSwitch := FALSE;
   BenchUut10.LeftLimitSwitch := FALSE;
   BenchUut10.RightLimitSwitch := FALSE;
   BenchUut10.GripLimitSwitch := FALSE;
   BenchUut10.ReleaseLimitSwitch := FALSE;
   TraceIn_ManualMode[87] := BenchUut10.ManualMode;
   TraceIn_SingleStepMode[87] := BenchUut10.SingleStepMode;
   TraceIn_SingleCycleMode[87] := BenchUut10.SingleCycleMode;
   TraceIn_ContinuousMode[87] := BenchUut10.ContinuousMode;
   TraceIn_EmergencyStop[87] := BenchUut10.EmergencyStop;
   TraceIn_Start[87] := BenchUut10.Start;
   TraceIn_DownButton[87] := BenchUut10.DownButton;
   TraceIn_UpButton[87] := BenchUut10.UpButton;
   TraceIn_LeftButton[87] := BenchUut10.LeftButton;
   TraceIn_RightButton[87] := BenchUut10.RightButton;
   TraceIn_GripButton[87] := BenchUut10.GripButton;
   TraceIn_ReleaseButton[87] := BenchUut10.ReleaseButton;
   TraceIn_DownLimitSwitch[87] := BenchUut10.DownLimitSwitch;
   TraceIn_UpLimitSwitch[87] := BenchUut10.UpLimitSwitch;
   TraceIn_LeftLimitSwitch[87] := BenchUut10.LeftLimitSwitch;
   TraceIn_RightLimitSwitch[87] := BenchUut10.RightLimitSwitch;
   TraceIn_GripLimitSwitch[87] := BenchUut10.GripLimitSwitch;
   TraceIn_ReleaseLimitSwitch[87] := BenchUut10.ReleaseLimitSwitch;
   BenchUut10();
   TraceOut_MoveDown[87] := BenchUut10.MoveDown;
   TraceOut_MoveUp[87] := BenchUut10.MoveUp;
   TraceOut_MoveLeft[87] := BenchUut10.MoveLeft;
   TraceOut_MoveRight[87] := BenchUut10.MoveRight;
   TraceOut_ActivateGrip[87] := BenchUut10.ActivateGrip;
   TraceOut_ActivateRelease[87] := BenchUut10.ActivateRelease;
   BenchCalls := BenchCalls + 1;
 88:
   BenchUut10.ManualMode := TRUE;
   BenchUut10.SingleStepMode := FALSE;
   BenchUut10.SingleCycleMode := FALSE;
   BenchUut10.ContinuousMode := FALSE;
   BenchUut10.EmergencyStop := TRUE;
   BenchUut10.Start := FALSE;
   BenchUut10.DownButton := FALSE;
   BenchUut10.UpButton := FALSE;
   BenchUut10.LeftButton := TRUE;
   BenchUut10.RightButton := FALSE;
   BenchUut10.GripButton := FALSE;
   BenchUut10.ReleaseButton := FALSE;
   BenchUut10.DownLimitSwitch := FALSE;
   BenchUut10.UpLimitSwitch := FALSE;
   BenchUut10.LeftLimitSwitch := FALSE;
   BenchUut10.RightLimitSwitch := FALSE;
   BenchUut10.GripLimitSwitch := FALSE;
   BenchUut10.ReleaseLimitSwitch := FALSE;
   TraceIn_ManualMode[88] := BenchUut10.ManualMode;
   TraceIn_SingleStepMode[88] := BenchUut10.SingleStepMode;
   TraceIn_SingleCycleMode[88] := BenchUut10.SingleCycleMode;
   TraceIn_ContinuousMode[88] := BenchUut10.ContinuousMode;
   TraceIn_EmergencyStop[88] := BenchUut10.EmergencyStop;
   TraceIn_Start[88] := BenchUut10.Start;
   TraceIn_DownButton[88] := BenchUut10.DownButton;
   TraceIn_UpButton[88] := BenchUut10.UpButton;
   TraceIn_LeftButton[88] := BenchUut10.LeftButton;
   TraceIn_RightButton[88] := BenchUut10.RightButton;
   TraceIn_GripButton[88] := BenchUut10.GripButton;
   TraceIn_ReleaseButton[88] := BenchUut10.ReleaseButton;
   TraceIn_DownLimitSwitch[88] := BenchUut10.DownLimitSwitch;
   TraceIn_UpLimitSwitch[88] := BenchUut10.UpLimitSwitch;
   TraceIn_LeftLimitSwitch[88] := BenchUut10.LeftLimitSwitch;
   TraceIn_RightLimitSwitch[88] := BenchUut10.RightLimitSwitch;
   TraceIn_GripLimitSwitch[88] := BenchUut10.GripLimitSwitch;
   TraceIn_ReleaseLimitSwitch[88] := BenchUut10.ReleaseLimitSwitch;
   BenchUut10();
   TraceOut_MoveDown[88] := BenchUut10.MoveDown;
   TraceOut_MoveUp[88] := BenchUut10.MoveUp;
   TraceOut_MoveLeft[88] := BenchUut10.MoveLeft;
   TraceOut_MoveRight[88] := BenchUut10.MoveRight;
   TraceOut_ActivateGrip[88] := BenchUut10.ActivateGrip;
   TraceOut_ActivateRelease[88] := BenchUut10.ActivateRelease;
   BenchCalls := BenchCalls + 1;
 89:
   BenchUut10.ManualMode := TRUE;
   BenchUut10.SingleStepMode := FALSE;
   BenchUut10.SingleCycleMode := FALSE;
   BenchUut10.ContinuousMode := FALSE;
   BenchUut10.EmergencyStop := TRUE;
   BenchUut10.Start := FALSE;
   BenchUut10.DownButton := FALSE;
   BenchUut10.UpButton := FALSE;
   BenchUut10.LeftButton := TRUE;
   BenchUut10.RightButton := FALSE;
   BenchUut10.GripButton := FALSE;
   BenchUut10.ReleaseButton := FALSE;
   BenchUut10.DownLimitSwitch := FALSE;
   BenchUut10.UpLimitSwitch := FALSE;
   BenchUut10.LeftLimitSwitch := FALSE;
   BenchUut10.RightLimitSwitch := FALSE;
   BenchUut10.GripLimitSwitch := FALSE;
   BenchUut10.ReleaseLimitSwitch := FALSE;
   TraceIn_ManualMode[89] := BenchUut10.ManualMode;
   TraceIn_SingleStepMode[89] := BenchUut10.SingleStepMode;
   TraceIn_SingleCycleMode[89] := BenchUut10.SingleCycleMode;
   TraceIn_ContinuousMode[89] := BenchUut10.ContinuousMode;
   TraceIn_EmergencyStop[89] := BenchUut10.EmergencyStop;
   TraceIn_Start[89] := BenchUut10.Start;
   TraceIn_DownButton[89] := BenchUut10.DownButton;
   TraceIn_UpButton[89] := BenchUut10.UpButton;
   TraceIn_LeftButton[89] := BenchUut10.LeftButton;
   TraceIn_RightButton[89] := BenchUut10.RightButton;
   TraceIn_GripButton[89] := BenchUut10.GripButton;
   TraceIn_ReleaseButton[89] := BenchUut10.ReleaseButton;
   TraceIn_DownLimitSwitch[89] := BenchUut10.DownLimitSwitch;
   TraceIn_UpLimitSwitch[89] := BenchUut10.UpLimitSwitch;
   TraceIn_LeftLimitSwitch[89] := BenchUut10.LeftLimitSwitch;
   TraceIn_RightLimitSwitch[89] := BenchUut10.RightLimitSwitch;
   TraceIn_GripLimitSwitch[89] := BenchUut10.GripLimitSwitch;
   TraceIn_ReleaseLimitSwitch[89] := BenchUut10.ReleaseLimitSwitch;
   BenchUut10();
   TraceOut_MoveDown[89] := BenchUut10.MoveDown;
   TraceOut_MoveUp[89] := BenchUut10.MoveUp;
   TraceOut_MoveLeft[89] := BenchUut10.MoveLeft;
   TraceOut_MoveRight[89] := BenchUut10.MoveRight;
   TraceOut_ActivateGrip[89] := BenchUut10.ActivateGrip;
   TraceOut_ActivateRelease[89] := BenchUut10.ActivateRelease;
   BenchCalls := BenchCalls + 1;
 90:
   BenchUut10.ManualMode := TRUE;
   BenchUut10.SingleStepMode := FALSE;
   BenchUut10.SingleCycleMode := FALSE;
   BenchUut10.ContinuousMode := FALSE;
   BenchUut10.EmergencyStop := TRUE;
   BenchUut10.Start := FALSE;
   BenchUut10.DownButton := FALSE;
   BenchUut10.UpButton := FALSE;
   BenchUut10.LeftButton := TRUE;
   BenchUut10.RightButton := FALSE;
   BenchUut10.GripButton := FALSE;
   BenchUut10.ReleaseButton := FALSE;
   BenchUut10.DownLimitSwitch := FALSE;
   BenchUut10.UpLimitSwitch := FALSE;
   BenchUut10.LeftLimitSwitch := TRUE;
   BenchUut10.RightLimitSwitch := FALSE;
   BenchUut10.GripLimitSwitch := FALSE;
   BenchUut10.ReleaseLimitSwitch := FALSE;
   TraceIn_ManualMode[90] := BenchUut10.ManualMode;
   TraceIn_SingleStepMode[90] := BenchUut10.SingleStepMode;
   TraceIn_SingleCycleMode[90] := BenchUut10.SingleCycleMode;
   TraceIn_ContinuousMode[90] := BenchUut10.ContinuousMode;
   TraceIn_EmergencyStop[90] := BenchUut10.EmergencyStop;
   TraceIn_Start[90] := BenchUut10.Start;
   TraceIn_DownButton[90] := BenchUut10.DownButton;
   TraceIn_UpButton[90] := BenchUut10.UpButton;
   TraceIn_LeftButton[90] := BenchUut10.LeftButton;
   TraceIn_RightButton[90] := BenchUut10.RightButton;
   TraceIn_GripButton[90] := BenchUut10.GripButton;
   TraceIn_ReleaseButton[90] := BenchUut10.ReleaseButton;
   TraceIn_DownLimitSwitch[90] := BenchUut10.DownLimitSwitch;
   TraceIn_UpLimitSwitch[90] := BenchUut10.UpLimitSwitch;
   TraceIn_LeftLimitSwitch[90] := BenchUut10.LeftLimitSwitch;
   TraceIn_RightLimitSwitch[90] := BenchUut10.RightLimitSwitch;
   TraceIn_GripLimitSwitch[90] := BenchUut10.GripLimitSwitch;
   TraceIn_ReleaseLimitSwitch[90] := BenchUut10.ReleaseLimitSwitch;
   BenchUut10();
   TraceOut_MoveDown[90] := BenchUut10.MoveDown;
   TraceOut_MoveUp[90] := BenchUut10.MoveUp;
   TraceOut_MoveLeft[90] := BenchUut10.MoveLeft;
   TraceOut_MoveRight[90] := BenchUut10.MoveRight;
   TraceOut_ActivateGrip[90] := BenchUut10.ActivateGrip;
   TraceOut_ActivateRelease[90] := BenchUut10.ActivateRelease;
   BenchCalls := BenchCalls + 1;
 91:
   BenchUut10.ManualMode := TRUE;
   BenchUut10.SingleStepMode := FALSE;
   BenchUut10.SingleCycleMode := FALSE;
   BenchUut10.ContinuousMode := FALSE;
   BenchUut10.EmergencyStop := TRUE;
   BenchUut10.Start := FALSE;
   BenchUut10.DownButton := FALSE;
   BenchUut10.UpButton := FALSE;
   BenchUut10.LeftButton := FALSE;
   BenchUut10.RightButton := FALSE;
   BenchUut10.GripButton := FALSE;
   BenchUut10.ReleaseButton := FALSE;
   BenchUut10.DownLimitSwitch := FALSE;
   BenchUut10.UpLimitSwitch := FALSE;
   BenchUut10.LeftLimitSwitch := TRUE;
   BenchUut10.RightLimitSwitch := FALSE;
   BenchUut10.GripLimitSwitch := FALSE;
   BenchUut10.ReleaseLimitSwitch := FALSE;
   TraceIn_ManualMode[91] := BenchUut10.ManualMode;
   TraceIn_SingleStepMode[91] := BenchUut10.SingleStepMode;
   TraceIn_SingleCycleMode[91] := BenchUut10.SingleCycleMode;
   TraceIn_ContinuousMode[91] := BenchUut10.ContinuousMode;
   TraceIn_EmergencyStop[91] := BenchUut10.EmergencyStop;
   TraceIn_Start[91] := BenchUut10.Start;
   TraceIn_DownButton[91] := BenchUut10.DownButton;
   TraceIn_UpButton[91] := BenchUut10.UpButton;
   TraceIn_LeftButton[91] := BenchUut10.LeftButton;
   TraceIn_RightButton[91] := BenchUut10.RightButton;
   TraceIn_GripButton[91] := BenchUut10.GripButton;
   TraceIn_ReleaseButton[91] := BenchUut10.ReleaseButton;
   TraceIn_DownLimitSwitch[91] := BenchUut10.DownLimitSwitch;
   TraceIn_UpLimitSwitch[91] := BenchUut10.UpLimitSwitch;
   TraceIn_LeftLimitSwitch[91] := BenchUut10.LeftLimitSwitch;
   TraceIn_RightLimitSwitch[91] := BenchUut10.RightLimitSwitch;
   TraceIn_GripLimitSwitch[91] := BenchUut10.GripLimitSwitch;
   TraceIn_ReleaseLimitSwitch[91] := BenchUut10.ReleaseLimitSwitch;
   BenchUut10();
   TraceOut_MoveDown[91] := BenchUut10.MoveDown;
   TraceOut_MoveUp[91] := BenchUut10.MoveUp;
   TraceOut_MoveLeft[91] := BenchUut10.MoveLeft;
   TraceOut_MoveRight[91] := BenchUut10.MoveRight;
   TraceOut_ActivateGrip[91] := BenchUut10.ActivateGrip;
   TraceOut_ActivateRelease[91] := BenchUut10.ActivateRelease;
   BenchCalls := BenchCalls + 1;
 92:
   BenchUut10.ManualMode := TRUE;
   BenchUut10.SingleStepMode := FALSE;
   BenchUut10.SingleCycleMode := FALSE;
   BenchUut10.ContinuousMode := FALSE;
   BenchUut10.EmergencyStop := TRUE;
   BenchUut10.Start := FALSE;
   BenchUut10.DownButton := FALSE;
   BenchUut10.UpButton := FALSE;
   BenchUut10.LeftButton := FALSE;
   BenchUut10.RightButton := FALSE;
   BenchUut10.GripButton := FALSE;
   BenchUut10.ReleaseButton := FALSE;
   BenchUut10.DownLimitSwitch := FALSE;
   BenchUut10.UpLimitSwitch := FALSE;
   BenchUut10.LeftLimitSwitch := FALSE;
   BenchUut10.RightLimitSwitch := FALSE;
   BenchUut10.GripLimitSwitch := FALSE;
   BenchUut10.ReleaseLimitSwitch := FALSE;
   TraceIn_ManualMode[92] := BenchUut10.ManualMode;
   TraceIn_SingleStepMode[92] := BenchUut10.SingleStepMode;
   TraceIn_SingleCycleMode[92] := BenchUut10.SingleCycleMode;
   TraceIn_ContinuousMode[92] := BenchUut10.ContinuousMode;
   TraceIn_EmergencyStop[92] := BenchUut10.EmergencyStop;
   TraceIn_Start[92] := BenchUut10.Start;
   TraceIn_DownButton[92] := BenchUut10.DownButton;
   TraceIn_UpButton[92] := BenchUut10.UpButton;
   TraceIn_LeftButton[92] := BenchUut10.LeftButton;
   TraceIn_RightButton[92] := BenchUut10.RightButton;
   TraceIn_GripButton[92] := BenchUut10.GripButton;
   TraceIn_ReleaseButton[92] := BenchUut10.ReleaseButton;
   TraceIn_DownLimitSwitch[92] := BenchUut10.DownLimitSwitch;
   TraceIn_UpLimitSwitch[92] := BenchUut10.UpLimitSwitch;
   TraceIn_LeftLimitSwitch[92] := BenchUut10.LeftLimitSwitch;
   TraceIn_RightLimitSwitch[92] := BenchUut10.RightLimitSwitch;
   TraceIn_GripLimitSwitch[92] := BenchUut10.GripLimitSwitch;
   TraceIn_ReleaseLimitSwitch[92] := BenchUut10.ReleaseLimitSwitch;
   BenchUut10();
   TraceOut_MoveDown[92] := BenchUut10.MoveDown;
   TraceOut_MoveUp[92] := BenchUut10.MoveUp;
   TraceOut_MoveLeft[92] := BenchUut10.MoveLeft;
   TraceOut_MoveRight[92] := BenchUut10.MoveRight;
   TraceOut_ActivateGrip[92] := BenchUut10.ActivateGrip;
   TraceOut_ActivateRelease[92] := BenchUut10.ActivateRelease;
   BenchCalls := BenchCalls + 1;
 93:
   BenchUut11.ManualMode := TRUE;
   BenchUut11.SingleStepMode := FALSE;
   BenchUut11.SingleCycleMode := FALSE;
   BenchUut11.ContinuousMode := FALSE;
   BenchUut11.EmergencyStop := TRUE;
   BenchUut11.Start := FALSE;
   BenchUut11.DownButton := FALSE;
   BenchUut11.UpButton := FALSE;
   BenchUut11.LeftButton := FALSE;
   BenchUut11.RightButton := FALSE;
   BenchUut11.GripButton := FALSE;
   BenchUut11.ReleaseButton := FALSE;
   BenchUut11.DownLimitSwitch := FALSE;
   BenchUut11.UpLimitSwitch := FALSE;
   BenchUut11.LeftLimitSwitch := FALSE;
   BenchUut11.RightLimitSwitch := FALSE;
   BenchUut11.GripLimitSwitch := FALSE;
   BenchUut11.ReleaseLimitSwitch := FALSE;
   TraceIn_ManualMode[93] := BenchUut11.ManualMode;
   TraceIn_SingleStepMode[93] := BenchUut11.SingleStepMode;
   TraceIn_SingleCycleMode[93] := BenchUut11.SingleCycleMode;
   TraceIn_ContinuousMode[93] := BenchUut11.ContinuousMode;
   TraceIn_EmergencyStop[93] := BenchUut11.EmergencyStop;
   TraceIn_Start[93] := BenchUut11.Start;
   TraceIn_DownButton[93] := BenchUut11.DownButton;
   TraceIn_UpButton[93] := BenchUut11.UpButton;
   TraceIn_LeftButton[93] := BenchUut11.LeftButton;
   TraceIn_RightButton[93] := BenchUut11.RightButton;
   TraceIn_GripButton[93] := BenchUut11.GripButton;
   TraceIn_ReleaseButton[93] := BenchUut11.ReleaseButton;
   TraceIn_DownLimitSwitch[93] := BenchUut11.DownLimitSwitch;
   TraceIn_UpLimitSwitch[93] := BenchUut11.UpLimitSwitch;
   TraceIn_LeftLimitSwitch[93] := BenchUut11.LeftLimitSwitch;
   TraceIn_RightLimitSwitch[93] := BenchUut11.RightLimitSwitch;
   TraceIn_GripLimitSwitch[93] := BenchUut11.GripLimitSwitch;
   TraceIn_ReleaseLimitSwitch[93] := BenchUut11.ReleaseLimitSwitch;
   BenchUut11();
   TraceOut_MoveDown[93] := BenchUut11.MoveDown;
   TraceOut_MoveUp[93] := BenchUut11.MoveUp;
   TraceOut_MoveLeft[93] := BenchUut11.MoveLeft;
   TraceOut_MoveRight[93] := BenchUut11.MoveRight;
   TraceOut_ActivateGrip[93] := BenchUut11.ActivateGrip;
   TraceOut_ActivateRelease[93] := BenchUut11.ActivateRelease;
   BenchCalls := BenchCalls + 1;
 94:
   BenchUut11.ManualMode := TRUE;
   BenchUut11.SingleStepMode := FALSE;
   BenchUut11.SingleCycleMode := FALSE;
   BenchUut11.ContinuousMode := FALSE;
   BenchUut11.EmergencyStop := TRUE;
   BenchUut11.Start := FALSE;
   BenchUut11.DownButton := FALSE;
   BenchUut11.UpButton := FALSE;
   BenchUut11.LeftButton := FALSE;
   BenchUut11.RightButton := TRUE;
   BenchUut11.GripButton := FALSE;
   BenchUut11.ReleaseButton := FALSE;
   BenchUut11.DownLimitSwitch := FALSE;
   BenchUut11.UpLimitSwitch := FALSE;
   BenchUut11.LeftLimitSwitch := FALSE;
   BenchUut11.RightLimitSwitch := FALSE;
   BenchUut11.GripLimitSwitch := FALSE;
   BenchUut11.ReleaseLimitSwitch := FALSE;
   TraceIn_ManualMode[94] := BenchUut11.ManualMode;
   TraceIn_SingleStepMode[94] := BenchUut11.SingleStepMode;
   TraceIn_SingleCycleMode[94] := BenchUut11.SingleCycleMode;
   TraceIn_ContinuousMode[94] := BenchUut11.ContinuousMode;
   TraceIn_EmergencyStop[94] := BenchUut11.EmergencyStop;
   TraceIn_Start[94] := BenchUut11.Start;
   TraceIn_DownButton[94] := BenchUut11.DownButton;
   TraceIn_UpButton[94] := BenchUut11.UpButton;
   TraceIn_LeftButton[94] := BenchUut11.LeftButton;
   TraceIn_RightButton[94] := BenchUut11.RightButton;
   TraceIn_GripButton[94] := BenchUut11.GripButton;
   TraceIn_ReleaseButton[94] := BenchUut11.ReleaseButton;
   TraceIn_DownLimitSwitch[94] := BenchUut11.DownLimitSwitch;
   TraceIn_UpLimitSwitch[94] := BenchUut11.UpLimitSwitch;
   TraceIn_LeftLimitSwitch[94] := BenchUut11.LeftLimitSwitch;
   TraceIn_RightLimitSwitch[94] := BenchUut11.RightLimitSwitch;
   TraceIn_GripLimitSwitch[94] := BenchUut11.GripLimitSwitch;
   TraceIn_ReleaseLimitSwitch[94] := BenchUut11.ReleaseLimitSwitch;
   BenchUut11();
   TraceOut_MoveDown[94] := BenchUut11.MoveDown;
   TraceOut_MoveUp[94] := BenchUut11.MoveUp;
   TraceOut_MoveLeft[94] := BenchUut11.MoveLeft;
   TraceOut_MoveRight[94] := BenchUut11.MoveRight;
   TraceOut_ActivateGrip[94] := BenchUut11.ActivateGrip;
   TraceOut_ActivateRelease[94] := BenchUut11.ActivateRelease;
   BenchCalls := BenchCalls + 1;
 95:
   BenchUut11.ManualMode := TRUE;
   BenchUut11.SingleStepMode := FALSE;
   BenchUut11.SingleCycleMode := FALSE;
   BenchUut11.ContinuousMode := FALSE;
   BenchUut11.EmergencyStop := TRUE;
   BenchUut11.Start := FALSE;
   BenchUut11.DownButton := FALSE;
   BenchUut11.UpButton := FALSE;
   BenchUut11.LeftButton := FALSE;
   BenchUut11.RightButton := TRUE;
   BenchUut11.GripButton := FALSE;
   BenchUut11.ReleaseButton := FALSE;
   BenchUut11.DownLimitSwitch := FALSE;
   BenchUut11.UpLimitSwitch := FALSE;
   BenchUut11.LeftLimitSwitch := FALSE;
   BenchUut11.RightLimitSwitch := FALSE;
   BenchUut11.GripLimitSwitch := FALSE;
   BenchUut11.ReleaseLimitSwitch := FALSE;
   TraceIn_ManualMode[95] := BenchUut11.ManualMode;
   TraceIn_SingleStepMode[95] := BenchUut11.SingleStepMode;
   TraceIn_SingleCycleMode[95] := BenchUut11.SingleCycleMode;
   TraceIn_ContinuousMode[95] := BenchUut11.ContinuousMode;
   TraceIn_EmergencyStop[95] := BenchUut11.EmergencyStop;
   TraceIn_Start[95] := BenchUut11.Start;
   TraceIn_DownButton[95] := BenchUut11.DownButton;
   TraceIn_UpButton[95] := BenchUut11.UpButton;
   TraceIn_LeftButton[95] := BenchUut11.LeftButton;
   TraceIn_RightButton[95] := BenchUut11.RightButton;
   TraceIn_GripButton[95] := BenchUut11.GripButton;
   TraceIn_ReleaseButton[95] := BenchUut11.ReleaseButton;
   TraceIn_DownLimitSwitch[95] := BenchUut11.DownLimitSwitch;
   TraceIn_UpLimitSwitch[95] := BenchUut11.UpLimitSwitch;
   TraceIn_LeftLimitSwitch[95] := BenchUut11.LeftLimitSwitch;
   TraceIn_RightLimitSwitch[95] := BenchUut11.RightLimitSwitch;
   TraceIn_GripLimitSwitch[95] := BenchUut11.GripLimitSwitch;
   TraceIn_ReleaseLimitSwitch[95] := BenchUut11.ReleaseLimitSwitch;
   BenchUut11();
   TraceOut_MoveDown[95] := BenchUut11.MoveDown;
   TraceOut_MoveUp[95] := BenchUut11.MoveUp;
   TraceOut_MoveLeft[95] := BenchUut11.MoveLeft;
   TraceOut_MoveRight[95] := BenchUut11.MoveRight;
   TraceOut_ActivateGrip[95] := BenchUut11.ActivateGrip;
   TraceOut_ActivateRelease[95] := BenchUut11.ActivateRelease;
   BenchCalls := BenchCalls + 1;
 96:
   BenchUut11.ManualMode := TRUE;
   BenchUut11.SingleStepMode := FALSE;
   BenchUut11.SingleCycleMode := FALSE;
   BenchUut11.ContinuousMode := FALSE;
   BenchUut11.EmergencyStop := TRUE;
   BenchUut11.Start := FALSE;
   BenchUut11.DownButton := FALSE;
   BenchUut11.UpButton := FALSE;
   BenchUut11.LeftButton := FALSE;
   BenchUut11.RightButton := TRUE;
   BenchUut11.GripButton := FALSE;
   BenchUut11.ReleaseButton := FALSE;
   BenchUut11.DownLimitSwitch := FALSE;
   BenchUut11.UpLimitSwitch := FALSE;
   BenchUut11.LeftLimitSwitch := FALSE;
   BenchUut11.RightLimitSwitch := TRUE;
   BenchUut11.GripLimitSwitch := FALSE;
   BenchUut11.ReleaseLimitSwitch := FALSE;
   TraceIn_ManualMode[96] := BenchUut11.ManualMode;
   TraceIn_SingleStepMode[96] := BenchUut11.SingleStepMode;
   TraceIn_SingleCycleMode[96] := BenchUut11.SingleCycleMode;
   TraceIn_ContinuousMode[96] := BenchUut11.ContinuousMode;
   TraceIn_EmergencyStop[96] := BenchUut11.EmergencyStop;
   TraceIn_Start[96] := BenchUut11.Start;
   TraceIn_DownButton[96] := BenchUut11.DownButton;
   TraceIn_UpButton[96] := BenchUut11.UpButton;
   TraceIn_LeftButton[96] := BenchUut11.LeftButton;
   TraceIn_RightButton[96] := BenchUut11.RightButton;
   TraceIn_GripButton[96] := BenchUut11.GripButton;
   TraceIn_ReleaseButton[96] := BenchUut11.ReleaseButton;
   TraceIn_DownLimitSwitch[96] := BenchUut11.DownLimitSwitch;
   TraceIn_UpLimitSwitch[96] := BenchUut11.UpLimitSwitch;
   TraceIn_LeftLimitSwitch[96] := BenchUut11.LeftLimitSwitch;
   TraceIn_RightLimitSwitch[96] := BenchUut11.RightLimitSwitch;
   TraceIn_GripLimitSwitch[96] := BenchUut11.GripLimitSwitch;
   TraceIn_ReleaseLimitSwitch[96] := BenchUut11.ReleaseLimitSwitch;
   BenchUut11();
   TraceOut_MoveDown[96] := BenchUut11.MoveDown;
   TraceOut_MoveUp[96] := BenchUut11.MoveUp;
   TraceOut_MoveLeft[96] := BenchUut11.MoveLeft;
   TraceOut_MoveRight[96] := BenchUut11.MoveRight;
   TraceOut_ActivateGrip[96] := BenchUut11.ActivateGrip;
   TraceOut_ActivateRelease[96] := BenchUut11.ActivateRelease;
   BenchCalls := BenchCalls + 1;
 97:
   BenchUut11.ManualMode := TRUE;
   BenchUut11.SingleStepMode := FALSE;
   BenchUut11.SingleCycleMode := FALSE;
   BenchUut11.ContinuousMode := FALSE;
   BenchUut11.EmergencyStop := TRUE;
   BenchUut11.Start := FALSE;
   BenchUut11.DownButton := FALSE;
   BenchUut11.UpButton := FALSE;
   BenchUut11.LeftButton := FALSE;
   BenchUut11.RightButton := FALSE;
   BenchUut11.GripButton := FALSE;
   BenchUut11.ReleaseButton := FALSE;
   BenchUut11.DownLimitSwitch := FALSE;
   BenchUut11.UpLimitSwitch := FALSE;
   BenchUut11.LeftLimitSwitch := FALSE;
   BenchUut11.RightLimitSwitch := TRUE;
   BenchUut11.GripLimitSwitch := FALSE;
   BenchUut11.ReleaseLimitSwitch := FALSE;
   TraceIn_ManualMode[97] := BenchUut11.ManualMode;
   TraceIn_SingleStepMode[97] := BenchUut11.SingleStepMode;
   TraceIn_SingleCycleMode[97] := BenchUut11.SingleCycleMode;
   TraceIn_ContinuousMode[97] := BenchUut11.ContinuousMode;
   TraceIn_EmergencyStop[97] := BenchUut11.EmergencyStop;
   TraceIn_Start[97] := BenchUut11.Start;
   TraceIn_DownButton[97] := BenchUut11.DownButton;
   TraceIn_UpButton[97] := BenchUut11.UpButton;
   TraceIn_LeftButton[97] := BenchUut11.LeftButton;
   TraceIn_RightButton[97] := BenchUut11.RightButton;
   TraceIn_GripButton[97] := BenchUut11.GripButton;
   TraceIn_ReleaseButton[97] := BenchUut11.ReleaseButton;
   TraceIn_DownLimitSwitch[97] := BenchUut11.DownLimitSwitch;
   TraceIn_UpLimitSwitch[97] := BenchUut11.UpLimitSwitch;
   TraceIn_LeftLimitSwitch[97] := BenchUut11.LeftLimitSwitch;
   TraceIn_RightLimitSwitch[97] := BenchUut11.RightLimitSwitch;
   TraceIn_GripLimitSwitch[97] := BenchUut11.GripLimitSwitch;
   TraceIn_ReleaseLimitSwitch[97] := BenchUut11.ReleaseLimitSwitch;
   BenchUut11();
   TraceOut_MoveDown[97] := BenchUut11.MoveDown;
   TraceOut_MoveUp[97] := BenchUut11.MoveUp;
   TraceOut_MoveLeft[97] := BenchUut11.MoveLeft;
   TraceOut_MoveRight[97] := BenchUut11.MoveRight;
   TraceOut_ActivateGrip[97] := BenchUut11.ActivateGrip;
   TraceOut_ActivateRelease[97] := BenchUut11.ActivateRelease;
   BenchCalls := BenchCalls + 1;
 98:
   BenchUut11.ManualMode := TRUE;
   BenchUut11.SingleStepMode := FALSE;
   BenchUut11.SingleCycleMode := FALSE;
   BenchUut11.ContinuousMode := FALSE;
   BenchUut11.EmergencyStop := TRUE;
   BenchUut11.Start := FALSE;
   BenchUut11.DownButton := FALSE;
   BenchUut11.UpButton := FALSE;
   BenchUut11.LeftButton := FALSE;
   BenchUut11.RightButton := FALSE;
   BenchUut11.GripButton := FALSE;
   BenchUut11.ReleaseButton := FALSE;
   BenchUut11.DownLimitSwitch := FALSE;
   BenchUut11.UpLimitSwitch := FALSE;
   BenchUut11.LeftLimitSwitch := FALSE;
   BenchUut11.RightLimitSwitch := FALSE;
   BenchUut11.GripLimitSwitch := FALSE;
   BenchUut11.ReleaseLimitSwitch := FALSE;
   TraceIn_ManualMode[98] := BenchUut11.ManualMode;
   TraceIn_SingleStepMode[98] := BenchUut11.SingleStepMode;
   TraceIn_SingleCycleMode[98] := BenchUut11.SingleCycleMode;
   TraceIn_ContinuousMode[98] := BenchUut11.ContinuousMode;
   TraceIn_EmergencyStop[98] := BenchUut11.EmergencyStop;
   TraceIn_Start[98] := BenchUut11.Start;
   TraceIn_DownButton[98] := BenchUut11.DownButton;
   TraceIn_UpButton[98] := BenchUut11.UpButton;
   TraceIn_LeftButton[98] := BenchUut11.LeftButton;
   TraceIn_RightButton[98] := BenchUut11.RightButton;
   TraceIn_GripButton[98] := BenchUut11.GripButton;
   TraceIn_ReleaseButton[98] := BenchUut11.ReleaseButton;
   TraceIn_DownLimitSwitch[98] := BenchUut11.DownLimitSwitch;
   TraceIn_UpLimitSwitch[98] := BenchUut11.UpLimitSwitch;
   TraceIn_LeftLimitSwitch[98] := BenchUut11.LeftLimitSwitch;
   TraceIn_RightLimitSwitch[98] := BenchUut11.RightLimitSwitch;
   TraceIn_GripLimitSwitch[98] := BenchUut11.GripLimitSwitch;
   TraceIn_ReleaseLimitSwitch[98] := BenchUut11.ReleaseLimitSwitch;
   BenchUut11();
   TraceOut_MoveDown[98] := BenchUut11.MoveDown;
   TraceOut_MoveUp[98] := BenchUut11.MoveUp;
   TraceOut_MoveLeft[98] := BenchUut11.MoveLeft;
   TraceOut_MoveRight[98] := BenchUut11.MoveRight;
   TraceOut_ActivateGrip[98] := BenchUut11.ActivateGrip;
   TraceOut_ActivateRelease[98] := BenchUut11.ActivateRelease;
   BenchCalls := BenchCalls + 1;
 99:
   BenchUut12.ManualMode := TRUE;
   BenchUut12.SingleStepMode := FALSE;
   BenchUut12.SingleCycleMode := FALSE;
   BenchUut12.ContinuousMode := FALSE;
   BenchUut12.EmergencyStop := TRUE;
   BenchUut12.Start := FALSE;
   BenchUut12.DownButton := FALSE;
   BenchUut12.UpButton := FALSE;
   BenchUut12.LeftButton := FALSE;
   BenchUut12.RightButton := FALSE;
   BenchUut12.GripButton := FALSE;
   BenchUut12.ReleaseButton := FALSE;
   BenchUut12.DownLimitSwitch := FALSE;
   BenchUut12.UpLimitSwitch := FALSE;
   BenchUut12.LeftLimitSwitch := FALSE;
   BenchUut12.RightLimitSwitch := FALSE;
   BenchUut12.GripLimitSwitch := FALSE;
   BenchUut12.ReleaseLimitSwitch := FALSE;
   TraceIn_ManualMode[99] := BenchUut12.ManualMode;
   TraceIn_SingleStepMode[99] := BenchUut12.SingleStepMode;
   TraceIn_SingleCycleMode[99] := BenchUut12.SingleCycleMode;
   TraceIn_ContinuousMode[99] := BenchUut12.ContinuousMode;
   TraceIn_EmergencyStop[99] := BenchUut12.EmergencyStop;
   TraceIn_Start[99] := BenchUut12.Start;
   TraceIn_DownButton[99] := BenchUut12.DownButton;
   TraceIn_UpButton[99] := BenchUut12.UpButton;
   TraceIn_LeftButton[99] := BenchUut12.LeftButton;
   TraceIn_RightButton[99] := BenchUut12.RightButton;
   TraceIn_GripButton[99] := BenchUut12.GripButton;
   TraceIn_ReleaseButton[99] := BenchUut12.ReleaseButton;
   TraceIn_DownLimitSwitch[99] := BenchUut12.DownLimitSwitch;
   TraceIn_UpLimitSwitch[99] := BenchUut12.UpLimitSwitch;
   TraceIn_LeftLimitSwitch[99] := BenchUut12.LeftLimitSwitch;
   TraceIn_RightLimitSwitch[99] := BenchUut12.RightLimitSwitch;
   TraceIn_GripLimitSwitch[99] := BenchUut12.GripLimitSwitch;
   TraceIn_ReleaseLimitSwitch[99] := BenchUut12.ReleaseLimitSwitch;
   BenchUut12();
   TraceOut_MoveDown[99] := BenchUut12.MoveDown;
   TraceOut_MoveUp[99] := BenchUut12.MoveUp;
   TraceOut_MoveLeft[99] := BenchUut12.MoveLeft;
   TraceOut_MoveRight[99] := BenchUut12.MoveRight;
   TraceOut_ActivateGrip[99] := BenchUut12.ActivateGrip;
   TraceOut_ActivateRelease[99] := BenchUut12.ActivateRelease;
   BenchCalls := BenchCalls + 1;
 100:
   BenchUut12.ManualMode := TRUE;
   BenchUut12.SingleStepMode := FALSE;
   BenchUut12.SingleCycleMode := FALSE;
   BenchUut12.ContinuousMode := FALSE;
   BenchUut12.EmergencyStop := TRUE;
   BenchUut12.Start := FALSE;
   BenchUut12.DownButton := FALSE;
   BenchUut12.UpButton := FALSE;
   BenchUut12.LeftButton := FALSE;
   BenchUut12.RightButton := FALSE;
   BenchUut12.GripButton := TRUE;
   BenchUut12.ReleaseButton := FALSE;
   BenchUut12.DownLimitSwitch := FALSE;
   BenchUut12.UpLimitSwitch := FALSE;
   BenchUut12.LeftLimitSwitch := FALSE;
   BenchUut12.RightLimitSwitch := FALSE;
   BenchUut12.GripLimitSwitch := FALSE;
   BenchUut12.ReleaseLimitSwitch := FALSE;
   TraceIn_ManualMode[100] := BenchUut12.ManualMode;
   TraceIn_SingleStepMode[100] := BenchUut12.SingleStepMode;
   TraceIn_SingleCycleMode[100] := BenchUut12.SingleCycleMode;
   TraceIn_ContinuousMode[100] := BenchUut12.ContinuousMode;
   TraceIn_EmergencyStop[100] := BenchUut12.EmergencyStop;
   TraceIn_Start[100] := BenchUut12.Start;
   TraceIn_DownButton[100] := BenchUut12.DownButton;
   TraceIn_UpButton[100] := BenchUut12.UpButton;
   TraceIn_LeftButton[100] := BenchUut12.LeftButton;
   TraceIn_RightButton[100] := BenchUut12.RightButton;
   TraceIn_GripButton[100] := BenchUut12.GripButton;
   TraceIn_ReleaseButton[100] := BenchUut12.ReleaseButton;
   TraceIn_DownLimitSwitch[100] := BenchUut12.DownLimitSwitch;
   TraceIn_UpLimitSwitch[100] := BenchUut12.UpLimitSwitch;
   TraceIn_LeftLimitSwitch[100] := BenchUut12.LeftLimitSwitch;
   TraceIn_RightLimitSwitch[100] := BenchUut12.RightLimitSwitch;
   TraceIn_GripLimitSwitch[100] := BenchUut12.GripLimitSwitch;
   TraceIn_ReleaseLimitSwitch[100] := BenchUut12.ReleaseLimitSwitch;
   BenchUut12();
   TraceOut_MoveDown[100] := BenchUut12.MoveDown;
   TraceOut_MoveUp[100] := BenchUut12.MoveUp;
   TraceOut_MoveLeft[100] := BenchUut12.MoveLeft;
   TraceOut_MoveRight[100] := BenchUut12.MoveRight;
   TraceOut_ActivateGrip[100] := BenchUut12.ActivateGrip;
   TraceOut_ActivateRelease[100] := BenchUut12.ActivateRelease;
   BenchCalls := BenchCalls + 1;
 101:
   BenchUut12.ManualMode := TRUE;
   BenchUut12.SingleStepMode := FALSE;
   BenchUut12.SingleCycleMode := FALSE;
   BenchUut12.ContinuousMode := FALSE;
   BenchUut12.EmergencyStop := TRUE;
   BenchUut12.Start := FALSE;
   BenchUut12.DownButton := FALSE;
   BenchUut12.UpButton := FALSE;
   BenchUut12.LeftButton := FALSE;
   BenchUut12.RightButton := FALSE;
   BenchUut12.GripButton := TRUE;
   BenchUut12.ReleaseButton := FALSE;
   BenchUut12.DownLimitSwitch := FALSE;
   BenchUut12.UpLimitSwitch := FALSE;
   BenchUut12.LeftLimitSwitch := FALSE;
   BenchUut12.RightLimitSwitch := FALSE;
   BenchUut12.GripLimitSwitch := FALSE;
   BenchUut12.ReleaseLimitSwitch := FALSE;
   TraceIn_ManualMode[101] := BenchUut12.ManualMode;
   TraceIn_SingleStepMode[101] := BenchUut12.SingleStepMode;
   TraceIn_SingleCycleMode[101] := BenchUut12.SingleCycleMode;
   TraceIn_ContinuousMode[101] := BenchUut12.ContinuousMode;
   TraceIn_EmergencyStop[101] := BenchUut12.EmergencyStop;
   TraceIn_Start[101] := BenchUut12.Start;
   TraceIn_DownButton[101] := BenchUut12.DownButton;
   TraceIn_UpButton[101] := BenchUut12.UpButton;
   TraceIn_LeftButton[101] := BenchUut12.LeftButton;
   TraceIn_RightButton[101] := BenchUut12.RightButton;
   TraceIn_GripButton[101] := BenchUut12.GripButton;
   TraceIn_ReleaseButton[101] := BenchUut12.ReleaseButton;
   TraceIn_DownLimitSwitch[101] := BenchUut12.DownLimitSwitch;
   TraceIn_UpLimitSwitch[101] := BenchUut12.UpLimitSwitch;
   TraceIn_LeftLimitSwitch[101] := BenchUut12.LeftLimitSwitch;
   TraceIn_RightLimitSwitch[101] := BenchUut12.RightLimitSwitch;
   TraceIn_GripLimitSwitch[101] := BenchUut12.GripLimitSwitch;
   TraceIn_ReleaseLimitSwitch[101] := BenchUut12.ReleaseLimitSwitch;
   BenchUut12();
   TraceOut_MoveDown[101] := BenchUut12.MoveDown;
   TraceOut_MoveUp[101] := BenchUut12.MoveUp;
   TraceOut_MoveLeft[101] := BenchUut12.MoveLeft;
   TraceOut_MoveRight[101] := BenchUut12.MoveRight;
   TraceOut_ActivateGrip[101] := BenchUut12.ActivateGrip;
   TraceOut_ActivateRelease[101] := BenchUut12.ActivateRelease;
   BenchCalls := BenchCalls + 1;
 102:
   BenchUut12.ManualMode := TRUE;
   BenchUut12.SingleStepMode := FALSE;
   BenchUut12.SingleCycleMode := FALSE;
   BenchUut12.ContinuousMode := FALSE;
   BenchUut12.EmergencyStop := TRUE;
   BenchUut12.Start := FALSE;
   BenchUut12.DownButton := FALSE;
   BenchUut12.UpButton := FALSE;
   BenchUut12.LeftButton := FALSE;
   BenchUut12.RightButton := FALSE;
   BenchUut12.GripButton := TRUE;
   BenchUut12.ReleaseButton := FALSE;
   BenchUut12.DownLimitSwitch := FALSE;
   BenchUut12.UpLimitSwitch := FALSE;
   BenchUut12.LeftLimitSwitch := FALSE;
   BenchUut12.RightLimitSwitch := FALSE;
   BenchUut12.GripLimitSwitch := TRUE;
   BenchUut12.ReleaseLimitSwitch := FALSE;
   TraceIn_ManualMode[102] := BenchUut12.ManualMode;
   TraceIn_SingleStepMode[102] := BenchUut12.SingleStepMode;
   TraceIn_SingleCycleMode[102] := BenchUut12.SingleCycleMode;
   TraceIn_ContinuousMode[102] := BenchUut12.ContinuousMode;
   TraceIn_EmergencyStop[102] := BenchUut12.EmergencyStop;
   TraceIn_Start[102] := BenchUut12.Start;
   TraceIn_DownButton[102] := BenchUut12.DownButton;
   TraceIn_UpButton[102] := BenchUut12.UpButton;
   TraceIn_LeftButton[102] := BenchUut12.LeftButton;
   TraceIn_RightButton[102] := BenchUut12.RightButton;
   TraceIn_GripButton[102] := BenchUut12.GripButton;
   TraceIn_ReleaseButton[102] := BenchUut12.ReleaseButton;
   TraceIn_DownLimitSwitch[102] := BenchUut12.DownLimitSwitch;
   TraceIn_UpLimitSwitch[102] := BenchUut12.UpLimitSwitch;
   TraceIn_LeftLimitSwitch[102] := BenchUut12.LeftLimitSwitch;
   TraceIn_RightLimitSwitch[102] := BenchUut12.RightLimitSwitch;
   TraceIn_GripLimitSwitch[102] := BenchUut12.GripLimitSwitch;
   TraceIn_ReleaseLimitSwitch[102] := BenchUut12.ReleaseLimitSwitch;
   BenchUut12();
   TraceOut_MoveDown[102] := BenchUut12.MoveDown;
   TraceOut_MoveUp[102] := BenchUut12.MoveUp;
   TraceOut_MoveLeft[102] := BenchUut12.MoveLeft;
   TraceOut_MoveRight[102] := BenchUut12.MoveRight;
   TraceOut_ActivateGrip[102] := BenchUut12.ActivateGrip;
   TraceOut_ActivateRelease[102] := BenchUut12.ActivateRelease;
   BenchCalls := BenchCalls + 1;
 103:
   BenchUut12.ManualMode := TRUE;
   BenchUut12.SingleStepMode := FALSE;
   BenchUut12.SingleCycleMode := FALSE;
   BenchUut12.ContinuousMode := FALSE;
   BenchUut12.EmergencyStop := TRUE;
   BenchUut12.Start := FALSE;
   BenchUut12.DownButton := FALSE;
   BenchUut12.UpButton := FALSE;
   BenchUut12.LeftButton := FALSE;
   BenchUut12.RightButton := FALSE;
   BenchUut12.GripButton := FALSE;
   BenchUut12.ReleaseButton := FALSE;
   BenchUut12.DownLimitSwitch := FALSE;
   BenchUut12.UpLimitSwitch := FALSE;
   BenchUut12.LeftLimitSwitch := FALSE;
   BenchUut12.RightLimitSwitch := FALSE;
   BenchUut12.GripLimitSwitch := TRUE;
   BenchUut12.ReleaseLimitSwitch := FALSE;
   TraceIn_ManualMode[103] := BenchUut12.ManualMode;
   TraceIn_SingleStepMode[103] := BenchUut12.SingleStepMode;
   TraceIn_SingleCycleMode[103] := BenchUut12.SingleCycleMode;
   TraceIn_ContinuousMode[103] := BenchUut12.ContinuousMode;
   TraceIn_EmergencyStop[103] := BenchUut12.EmergencyStop;
   TraceIn_Start[103] := BenchUut12.Start;
   TraceIn_DownButton[103] := BenchUut12.DownButton;
   TraceIn_UpButton[103] := BenchUut12.UpButton;
   TraceIn_LeftButton[103] := BenchUut12.LeftButton;
   TraceIn_RightButton[103] := BenchUut12.RightButton;
   TraceIn_GripButton[103] := BenchUut12.GripButton;
   TraceIn_ReleaseButton[103] := BenchUut12.ReleaseButton;
   TraceIn_DownLimitSwitch[103] := BenchUut12.DownLimitSwitch;
   TraceIn_UpLimitSwitch[103] := BenchUut12.UpLimitSwitch;
   TraceIn_LeftLimitSwitch[103] := BenchUut12.LeftLimitSwitch;
   TraceIn_RightLimitSwitch[103] := BenchUut12.RightLimitSwitch;
   TraceIn_GripLimitSwitch[103] := BenchUut12.GripLimitSwitch;
   TraceIn_ReleaseLimitSwitch[103] := BenchUut12.ReleaseLimitSwitch;
   BenchUut12();
   TraceOut_MoveDown[103] := BenchUut12.MoveDown;
   TraceOut_MoveUp[103] := BenchUut12.MoveUp;
   TraceOut_MoveLeft[103] := BenchUut12.MoveLeft;
   TraceOut_MoveRight[103] := BenchUut12.MoveRight;
   TraceOut_ActivateGrip[103] := BenchUut12.ActivateGrip;
   TraceOut_ActivateRelease[103] := BenchUut12.ActivateRelease;
   BenchCalls := BenchCalls + 1;
 104:
   BenchUut12.ManualMode := TRUE;
   BenchUut12.SingleStepMode := FALSE;
   BenchUut12.SingleCycleMode := FALSE;
   BenchUut12.ContinuousMode := FALSE;
   BenchUut12.EmergencyStop := TRUE;
   BenchUut12.Start := FALSE;
   BenchUut12.DownButton := FALSE;
   BenchUut12.UpButton := FALSE;
   BenchUut12.LeftButton := FALSE;
   BenchUut12.RightButton := FALSE;
   BenchUut12.GripButton := FALSE;
   BenchUut12.ReleaseButton := FALSE;
   BenchUut12.DownLimitSwitch := FALSE;
   BenchUut12.UpLimitSwitch := FALSE;
   BenchUut12.LeftLimitSwitch := FALSE;
   BenchUut12.RightLimitSwitch := FALSE;
   BenchUut12.GripLimitSwitch := FALSE;
   BenchUut12.ReleaseLimitSwitch := FALSE;
   TraceIn_ManualMode[104] := BenchUut12.ManualMode;
   TraceIn_SingleStepMode[104] := BenchUut12.SingleStepMode;
   TraceIn_SingleCycleMode[104] := BenchUut12.SingleCycleMode;
   TraceIn_ContinuousMode[104] := BenchUut12.ContinuousMode;
   TraceIn_EmergencyStop[104] := BenchUut12.EmergencyStop;
   TraceIn_Start[104] := BenchUut12.Start;
   TraceIn_DownButton[104] := BenchUut12.DownButton;
   TraceIn_UpButton[104] := BenchUut12.UpButton;
   TraceIn_LeftButton[104] := BenchUut12.LeftButton;
   TraceIn_RightButton[104] := BenchUut12.RightButton;
   TraceIn_GripButton[104] := BenchUut12.GripButton;
   TraceIn_ReleaseButton[104] := BenchUut12.ReleaseButton;
   TraceIn_DownLimitSwitch[104] := BenchUut12.DownLimitSwitch;
   TraceIn_UpLimitSwitch[104] := BenchUut12.UpLimitSwitch;
   TraceIn_LeftLimitSwitch[104] := BenchUut12.LeftLimitSwitch;
   TraceIn_RightLimitSwitch[104] := BenchUut12.RightLimitSwitch;
   TraceIn_GripLimitSwitch[104] := BenchUut12.GripLimitSwitch;
   TraceIn_ReleaseLimitSwitch[104] := BenchUut12.ReleaseLimitSwitch;
   BenchUut12();
   TraceOut_MoveDown[104] := BenchUut12.MoveDown;
   TraceOut_MoveUp[104] := BenchUut12.MoveUp;
   TraceOut_MoveLeft[104] := BenchUut12.MoveLeft;
   TraceOut_MoveRight[104] := BenchUut12.MoveRight;
   TraceOut_ActivateGrip[104] := BenchUut12.ActivateGrip;
   TraceOut_ActivateRelease[104] := BenchUut12.ActivateRelease;
   BenchCalls := BenchCalls + 1;
 105:
   BenchUut13.ManualMode := TRUE;
   BenchUut13.SingleStepMode := FALSE;
   BenchUut13.SingleCycleMode := FALSE;
   BenchUut13.ContinuousMode := FALSE;
   BenchUut13.EmergencyStop := TRUE;
   BenchUut13.Start := FALSE;
   BenchUut13.DownButton := FALSE;
   BenchUut13.UpButton := FALSE;
   BenchUut13.LeftButton := FALSE;
   BenchUut13.RightButton := FALSE;
   BenchUut13.GripButton := FALSE;
   BenchUut13.ReleaseButton := FALSE;
   BenchUut13.DownLimitSwitch := FALSE;
   BenchUut13.UpLimitSwitch := FALSE;
   BenchUut13.LeftLimitSwitch := FALSE;
   BenchUut13.RightLimitSwitch := FALSE;
   BenchUut13.GripLimitSwitch := FALSE;
   BenchUut13.ReleaseLimitSwitch := FALSE;
   TraceIn_ManualMode[105] := BenchUut13.ManualMode;
   TraceIn_SingleStepMode[105] := BenchUut13.SingleStepMode;
   TraceIn_SingleCycleMode[105] := BenchUut13.SingleCycleMode;
   TraceIn_ContinuousMode[105] := BenchUut13.ContinuousMode;
   TraceIn_EmergencyStop[105] := BenchUut13.EmergencyStop;
   TraceIn_Start[105] := BenchUut13.Start;
   TraceIn_DownButton[105] := BenchUut13.DownButton;
   TraceIn_UpButton[105] := BenchUut13.UpButton;
   TraceIn_LeftButton[105] := BenchUut13.LeftButton;
   TraceIn_RightButton[105] := BenchUut13.RightButton;
   TraceIn_GripButton[105] := BenchUut13.GripButton;
   TraceIn_ReleaseButton[105] := BenchUut13.ReleaseButton;
   TraceIn_DownLimitSwitch[105] := BenchUut13.DownLimitSwitch;
   TraceIn_UpLimitSwitch[105] := BenchUut13.UpLimitSwitch;
   TraceIn_LeftLimitSwitch[105] := BenchUut13.LeftLimitSwitch;
   TraceIn_RightLimitSwitch[105] := BenchUut13.RightLimitSwitch;
   TraceIn_GripLimitSwitch[105] := BenchUut13.GripLimitSwitch;
   TraceIn_ReleaseLimitSwitch[105] := BenchUut13.ReleaseLimitSwitch;
   BenchUut13();
   TraceOut_MoveDown[105] := BenchUut13.MoveDown;
   TraceOut_MoveUp[105] := BenchUut13.MoveUp;
   TraceOut_MoveLeft[105] := BenchUut13.MoveLeft;
   TraceOut_MoveRight[105] := BenchUut13.MoveRight;
   TraceOut_ActivateGrip[105] := BenchUut13.ActivateGrip;
   TraceOut_ActivateRelease[105] := BenchUut13.ActivateRelease;
   BenchCalls := BenchCalls + 1;
 106:
   BenchUut13.ManualMode := TRUE;
   BenchUut13.SingleStepMode := FALSE;
   BenchUut13.SingleCycleMode := FALSE;
   BenchUut13.ContinuousMode := FALSE;
   BenchUut13.EmergencyStop := TRUE;
   BenchUut13.Start := FALSE;
   BenchUut13.DownButton := FALSE;
   BenchUut13.UpButton := FALSE;
   BenchUut13.LeftButton := FALSE;
   BenchUut13.RightButton := FALSE;
   BenchUut13.GripButton := FALSE;
   BenchUut13.ReleaseButton := TRUE;
   BenchUut13.DownLimitSwitch := FALSE;
   BenchUut13.UpLimitSwitch := FALSE;
   BenchUut13.LeftLimitSwitch := FALSE;
   BenchUut13.RightLimitSwitch := FALSE;
   BenchUut13.GripLimitSwitch := FALSE;
   BenchUut13.ReleaseLimitSwitch := FALSE;
   TraceIn_ManualMode[106] := BenchUut13.ManualMode;
   TraceIn_SingleStepMode[106] := BenchUut13.SingleStepMode;
   TraceIn_SingleCycleMode[106] := BenchUut13.SingleCycleMode;
   TraceIn_ContinuousMode[106] := BenchUut13.ContinuousMode;
   TraceIn_EmergencyStop[106] := BenchUut13.EmergencyStop;
   TraceIn_Start[106] := BenchUut13.Start;
   TraceIn_DownButton[106] := BenchUut13.DownButton;
   TraceIn_UpButton[106] := BenchUut13.UpButton;
   TraceIn_LeftButton[106] := BenchUut13.LeftButton;
   TraceIn_RightButton[106] := BenchUut13.RightButton;
   TraceIn_GripButton[106] := BenchUut13.GripButton;
   TraceIn_ReleaseButton[106] := BenchUut13.ReleaseButton;
   TraceIn_DownLimitSwitch[106] := BenchUut13.DownLimitSwitch;
   TraceIn_UpLimitSwitch[106] := BenchUut13.UpLimitSwitch;
   TraceIn_LeftLimitSwitch[106] := BenchUut13.LeftLimitSwitch;
   TraceIn_RightLimitSwitch[106] := BenchUut13.RightLimitSwitch;
   TraceIn_GripLimitSwitch[106] := BenchUut13.GripLimitSwitch;
   TraceIn_ReleaseLimitSwitch[106] := BenchUut13.ReleaseLimitSwitch;
   BenchUut13();
   TraceOut_MoveDown[106] := BenchUut13.MoveDown;
   TraceOut_MoveUp[106] := BenchUut13.MoveUp;
   TraceOut_MoveLeft[106] := BenchUut13.MoveLeft;
   TraceOut_MoveRight[106] := BenchUut13.MoveRight;
   TraceOut_ActivateGrip[106] := BenchUut13.ActivateGrip;
   TraceOut_ActivateRelease[106] := BenchUut13.ActivateRelease;
   BenchCalls := BenchCalls + 1;
 107:
   BenchUut13.ManualMode := TRUE;
   BenchUut13.SingleStepMode := FALSE;
   BenchUut13.SingleCycleMode := FALSE;
   BenchUut13.ContinuousMode := FALSE;
   BenchUut13.EmergencyStop := TRUE;
   BenchUut13.Start := FALSE;
   BenchUut13.DownButton := FALSE;
   BenchUut13.UpButton := FALSE;
   BenchUut13.LeftButton := FALSE;
   BenchUut13.RightButton := FALSE;
   BenchUut13.GripButton := FALSE;
   BenchUut13.ReleaseButton := TRUE;
   BenchUut13.DownLimitSwitch := FALSE;
   BenchUut13.UpLimitSwitch := FALSE;
   BenchUut13.LeftLimitSwitch := FALSE;
   BenchUut13.RightLimitSwitch := FALSE;
   BenchUut13.GripLimitSwitch := FALSE;
   BenchUut13.ReleaseLimitSwitch := FALSE;
   TraceIn_ManualMode[107] := BenchUut13.ManualMode;
   TraceIn_SingleStepMode[107] := BenchUut13.SingleStepMode;
   TraceIn_SingleCycleMode[107] := BenchUut13.SingleCycleMode;
   TraceIn_ContinuousMode[107] := BenchUut13.ContinuousMode;
   TraceIn_EmergencyStop[107] := BenchUut13.EmergencyStop;
   TraceIn_Start[107] := BenchUut13.Start;
   TraceIn_DownButton[107] := BenchUut13.DownButton;
   TraceIn_UpButton[107] := BenchUut13.UpButton;
   TraceIn_LeftButton[107] := BenchUut13.LeftButton;
   TraceIn_RightButton[107] := BenchUut13.RightButton;
   TraceIn_GripButton[107] := BenchUut13.GripButton;
   TraceIn_ReleaseButton[107] := BenchUut13.ReleaseButton;
   TraceIn_DownLimitSwitch[107] := BenchUut13.DownLimitSwitch;
   TraceIn_UpLimitSwitch[107] := BenchUut13.UpLimitSwitch;
   TraceIn_LeftLimitSwitch[107] := BenchUut13.LeftLimitSwitch;
   TraceIn_RightLimitSwitch[107] := BenchUut13.RightLimitSwitch;
   TraceIn_GripLimitSwitch[107] := BenchUut13.GripLimitSwitch;
   TraceIn_ReleaseLimitSwitch[107] := BenchUut13.ReleaseLimitSwitch;
   BenchUut13();
   TraceOut_MoveDown[107] := BenchUut13.MoveDown;
   TraceOut_MoveUp[107] := BenchUut13.MoveUp;
   TraceOut_MoveLeft[107] := BenchUut13.MoveLeft;
   TraceOut_MoveRight[107] := BenchUut13.MoveRight;
   TraceOut_ActivateGrip[107] := BenchUut13.ActivateGrip;
   TraceOut_ActivateRelease[107] := BenchUut13.ActivateRelease;
   BenchCalls := BenchCalls + 1;
 108:
   BenchUut13.ManualMode := TRUE;
   BenchUut13.SingleStepMode := FALSE;
   BenchUut13.SingleCycleMode := FALSE;
   BenchUut13.ContinuousMode := FALSE;
   BenchUut13.EmergencyStop := TRUE;
   BenchUut13.Start := FALSE;
   BenchUut13.DownButton := FALSE;
   BenchUut13.UpButton := FALSE;
   BenchUut13.LeftButton := FALSE;
   BenchUut13.RightButton := FALSE;
   BenchUut13.GripButton := FALSE;
   BenchUut13.ReleaseButton := TRUE;
   BenchUut13.DownLimitSwitch := FALSE;
   BenchUut13.UpLimitSwitch := FALSE;
   BenchUut13.LeftLimitSwitch := FALSE;
   BenchUut13.RightLimitSwitch := FALSE;
   BenchUut13.GripLimitSwitch := FALSE;
   BenchUut13.ReleaseLimitSwitch := TRUE;
   TraceIn_ManualMode[108] := BenchUut13.ManualMode;
   TraceIn_SingleStepMode[108] := BenchUut13.SingleStepMode;
   TraceIn_SingleCycleMode[108] := BenchUut13.SingleCycleMode;
   TraceIn_ContinuousMode[108] := BenchUut13.ContinuousMode;
   TraceIn_EmergencyStop[108] := BenchUut13.EmergencyStop;
   TraceIn_Start[108] := BenchUut13.Start;
   TraceIn_DownButton[108] := BenchUut13.DownButton;
   TraceIn_UpButton[108] := BenchUut13.UpButton;
   TraceIn_LeftButton[108] := BenchUut13.LeftButton;
   TraceIn_RightButton[108] := BenchUut13.RightButton;
   TraceIn_GripButton[108] := BenchUut13.GripButton;
   TraceIn_ReleaseButton[108] := BenchUut13.ReleaseButton;
   TraceIn_DownLimitSwitch[108] := BenchUut13.DownLimitSwitch;
   TraceIn_UpLimitSwitch[108] := BenchUut13.UpLimitSwitch;
   TraceIn_LeftLimitSwitch[108] := BenchUut13.LeftLimitSwitch;
   TraceIn_RightLimitSwitch[108] := BenchUut13.RightLimitSwitch;
   TraceIn_GripLimitSwitch[108] := BenchUut13.GripLimitSwitch;
   TraceIn_ReleaseLimitSwitch[108] := BenchUut13.ReleaseLimitSwitch;
   BenchUut13();
   TraceOut_MoveDown[108] := BenchUut13.MoveDown;
   TraceOut_MoveUp[108] := BenchUut13.MoveUp;
   TraceOut_MoveLeft[108] := BenchUut13.MoveLeft;
   TraceOut_MoveRight[108] := BenchUut13.MoveRight;
   TraceOut_ActivateGrip[108] := BenchUut13.ActivateGrip;
   TraceOut_ActivateRelease[108] := BenchUut13.ActivateRelease;
   BenchCalls := BenchCalls + 1;
 109:
   BenchUut13.ManualMode := TRUE;
   BenchUut13.SingleStepMode := FALSE;
   BenchUut13.SingleCycleMode := FALSE;
   BenchUut13.ContinuousMode := FALSE;
   BenchUut13.EmergencyStop := TRUE;
   BenchUut13.Start := FALSE;
   BenchUut13.DownButton := FALSE;
   BenchUut13.UpButton := FALSE;
   BenchUut13.LeftButton := FALSE;
   BenchUut13.RightButton := FALSE;
   BenchUut13.GripButton := FALSE;
   BenchUut13.ReleaseButton := FALSE;
   BenchUut13.DownLimitSwitch := FALSE;
   BenchUut13.UpLimitSwitch := FALSE;
   BenchUut13.LeftLimitSwitch := FALSE;
   BenchUut13.RightLimitSwitch := FALSE;
   BenchUut13.GripLimitSwitch := FALSE;
   BenchUut13.ReleaseLimitSwitch := TRUE;
   TraceIn_ManualMode[109] := BenchUut13.ManualMode;
   TraceIn_SingleStepMode[109] := BenchUut13.SingleStepMode;
   TraceIn_SingleCycleMode[109] := BenchUut13.SingleCycleMode;
   TraceIn_ContinuousMode[109] := BenchUut13.ContinuousMode;
   TraceIn_EmergencyStop[109] := BenchUut13.EmergencyStop;
   TraceIn_Start[109] := BenchUut13.Start;
   TraceIn_DownButton[109] := BenchUut13.DownButton;
   TraceIn_UpButton[109] := BenchUut13.UpButton;
   TraceIn_LeftButton[109] := BenchUut13.LeftButton;
   TraceIn_RightButton[109] := BenchUut13.RightButton;
   TraceIn_GripButton[109] := BenchUut13.GripButton;
   TraceIn_ReleaseButton[109] := BenchUut13.ReleaseButton;
   TraceIn_DownLimitSwitch[109] := BenchUut13.DownLimitSwitch;
   TraceIn_UpLimitSwitch[109] := BenchUut13.UpLimitSwitch;
   TraceIn_LeftLimitSwitch[109] := BenchUut13.LeftLimitSwitch;
   TraceIn_RightLimitSwitch[109] := BenchUut13.RightLimitSwitch;
   TraceIn_GripLimitSwitch[109] := BenchUut13.GripLimitSwitch;
   TraceIn_ReleaseLimitSwitch[109] := BenchUut13.ReleaseLimitSwitch;
   BenchUut13();
   TraceOut_MoveDown[109] := BenchUut13.MoveDown;
   TraceOut_MoveUp[109] := BenchUut13.MoveUp;
   TraceOut_MoveLeft[109] := BenchUut13.MoveLeft;
   TraceOut_MoveRight[109] := BenchUut13.MoveRight;
   TraceOut_ActivateGrip[109] := BenchUut13.ActivateGrip;
   TraceOut_ActivateRelease[109] := BenchUut13.ActivateRelease;
   BenchCalls := BenchCalls + 1;
 110:
   BenchUut13.ManualMode := TRUE;
   BenchUut13.SingleStepMode := FALSE;
   BenchUut13.SingleCycleMode := FALSE;
   BenchUut13.ContinuousMode := FALSE;
   BenchUut13.EmergencyStop := TRUE;
   BenchUut13.Start := FALSE;
   BenchUut13.DownButton := FALSE;
   BenchUut13.UpButton := FALSE;
   BenchUut13.LeftButton := FALSE;
   BenchUut13.RightButton := FALSE;
   BenchUut13.GripButton := FALSE;
   BenchUut13.ReleaseButton := FALSE;
   BenchUut13.DownLimitSwitch := FALSE;
   BenchUut13.UpLimitSwitch := FALSE;
   BenchUut13.LeftLimitSwitch := FALSE;
   BenchUut13.RightLimitSwitch := FALSE;
   BenchUut13.GripLimitSwitch := FALSE;
   BenchUut13.ReleaseLimitSwitch := FALSE;
   TraceIn_ManualMode[110] := BenchUut13.ManualMode;
   TraceIn_SingleStepMode[110] := BenchUut13.SingleStepMode;
   TraceIn_SingleCycleMode[110] := BenchUut13.SingleCycleMode;
   TraceIn_ContinuousMode[110] := BenchUut13.ContinuousMode;
   TraceIn_EmergencyStop[110] := BenchUut13.EmergencyStop;
   TraceIn_Start[110] := BenchUut13.Start;
   TraceIn_DownButton[110] := BenchUut13.DownButton;
   TraceIn_UpButton[110] := BenchUut13.UpButton;
   TraceIn_LeftButton[110] := BenchUut13.LeftButton;
   TraceIn_RightButton[110] := BenchUut13.RightButton;
   TraceIn_GripButton[110] := BenchUut13.GripButton;
   TraceIn_ReleaseButton[110] := BenchUut13.ReleaseButton;
   TraceIn_DownLimitSwitch[110] := BenchUut13.DownLimitSwitch;
   TraceIn_UpLimitSwitch[110] := BenchUut13.UpLimitSwitch;
   TraceIn_LeftLimitSwitch[110] := BenchUut13.LeftLimitSwitch;
   TraceIn_RightLimitSwitch[110] := BenchUut13.RightLimitSwitch;
   TraceIn_GripLimitSwitch[110] := BenchUut13.GripLimitSwitch;
   TraceIn_ReleaseLimitSwitch[110] := BenchUut13.ReleaseLimitSwitch;
   BenchUut13();
   TraceOut_MoveDown[110] := BenchUut13.MoveDown;
   TraceOut_MoveUp[110] := BenchUut13.MoveUp;
   TraceOut_MoveLeft[110] := BenchUut13.MoveLeft;
   TraceOut_MoveRight[110] := BenchUut13.MoveRight;
   TraceOut_ActivateGrip[110] := BenchUut13.ActivateGrip;
   TraceOut_ActivateRelease[110] := BenchUut13.ActivateRelease;
   BenchCalls := BenchCalls + 1;
 111:
   BenchUut14.ManualMode := FALSE;
   BenchUut14.SingleStepMode := TRUE;
   BenchUut14.SingleCycleMode := FALSE;
   BenchUut14.ContinuousMode := FALSE;
   BenchUut14.EmergencyStop := TRUE;
   BenchUut14.Start := FALSE;
   BenchUut14.DownButton := FALSE;
   BenchUut14.UpButton := FALSE;
   BenchUut14.LeftButton := FALSE;
   BenchUut14.RightButton := FALSE;
   BenchUut14.GripButton := FALSE;
   BenchUut14.ReleaseButton := FALSE;
   BenchUut14.DownLimitSwitch := FALSE;
   BenchUut14.UpLimitSwitch := TRUE;
   BenchUut14.LeftLimitSwitch := TRUE;
   BenchUut14.RightLimitSwitch := FALSE;
   BenchUut14.GripLimitSwitch := FALSE;
   BenchUut14.ReleaseLimitSwitch := FALSE;
   TraceIn_ManualMode[111] := BenchUut14.ManualMode;
   TraceIn_SingleStepMode[111] := BenchUut14.SingleStepMode;
   TraceIn_SingleCycleMode[111] := BenchUut14.SingleCycleMode;
   TraceIn_ContinuousMode[111] := BenchUut14.ContinuousMode;
   TraceIn_EmergencyStop[111] := BenchUut14.EmergencyStop;
   TraceIn_Start[111] := BenchUut14.Start;
   TraceIn_DownButton[111] := BenchUut14.DownButton;
   TraceIn_UpButton[111] := BenchUut14.UpButton;
   TraceIn_LeftButton[111] := BenchUut14.LeftButton;
   TraceIn_RightButton[111] := BenchUut14.RightButton;
   TraceIn_GripButton[111] := BenchUut14.GripButton;
   TraceIn_ReleaseButton[111] := BenchUut14.ReleaseButton;
   TraceIn_DownLimitSwitch[111] := BenchUut14.DownLimitSwitch;
   TraceIn_UpLimitSwitch[111] := BenchUut14.UpLimitSwitch;
   TraceIn_LeftLimitSwitch[111] := BenchUut14.LeftLimitSwitch;
   TraceIn_RightLimitSwitch[111] := BenchUut14.RightLimitSwitch;
   TraceIn_GripLimitSwitch[111] := BenchUut14.GripLimitSwitch;
   TraceIn_ReleaseLimitSwitch[111] := BenchUut14.ReleaseLimitSwitch;
   BenchUut14();
   TraceOut_MoveDown[111] := BenchUut14.MoveDown;
   TraceOut_MoveUp[111] := BenchUut14.MoveUp;
   TraceOut_MoveLeft[111] := BenchUut14.MoveLeft;
   TraceOut_MoveRight[111] := BenchUut14.MoveRight;
   TraceOut_ActivateGrip[111] := BenchUut14.ActivateGrip;
   TraceOut_ActivateRelease[111] := BenchUut14.ActivateRelease;
   BenchCalls := BenchCalls + 1;
 112:
   BenchUut14.ManualMode := FALSE;
   BenchUut14.SingleStepMode := TRUE;
   BenchUut14.SingleCycleMode := FALSE;
   BenchUut14.ContinuousMode := FALSE;
   BenchUut14.EmergencyStop := TRUE;
   BenchUut14.Start := TRUE;
   BenchUut14.DownButton := FALSE;
   BenchUut14.UpButton := FALSE;
   BenchUut14.LeftButton := FALSE;
   BenchUut14.RightButton := FALSE;
   BenchUut14.GripButton := FALSE;
   BenchUut14.ReleaseButton := FALSE;
   BenchUut14.DownLimitSwitch := FALSE;
   BenchUut14.UpLimitSwitch := TRUE;
   BenchUut14.LeftLimitSwitch := TRUE;
   BenchUut14.RightLimitSwitch := FALSE;
   BenchUut14.GripLimitSwitch := FALSE;
   BenchUut14.ReleaseLimitSwitch := FALSE;
   TraceIn_ManualMode[112] := BenchUut14.ManualMode;
   TraceIn_SingleStepMode[112] := BenchUut14.SingleStepMode;
   TraceIn_SingleCycleMode[112] := BenchUut14.SingleCycleMode;
   TraceIn_ContinuousMode[112] := BenchUut14.ContinuousMode;
   TraceIn_EmergencyStop[112] := BenchUut14.EmergencyStop;
   TraceIn_Start[112] := BenchUut14.Start;
   TraceIn_DownButton[112] := BenchUut14.DownButton;
   TraceIn_UpButton[112] := BenchUut14.UpButton;
   TraceIn_LeftButton[112] := BenchUut14.LeftButton;
   TraceIn_RightButton[112] := BenchUut14.RightButton;
   TraceIn_GripButton[112] := BenchUut14.GripButton;
   TraceIn_ReleaseButton[112] := BenchUut14.ReleaseButton;
   TraceIn_DownLimitSwitch[112] := BenchUut14.DownLimitSwitch;
   TraceIn_UpLimitSwitch[112] := BenchUut14.UpLimitSwitch;
   TraceIn_LeftLimitSwitch[112] := BenchUut14.LeftLimitSwitch;
   TraceIn_RightLimitSwitch[112] := BenchUut14.RightLimitSwitch;
   TraceIn_GripLimitSwitch[112] := BenchUut14.GripLimitSwitch;
   TraceIn_ReleaseLimitSwitch[112] := BenchUut14.ReleaseLimitSwitch;
   BenchUut14();
   TraceOut_MoveDown[112] := BenchUut14.MoveDown;
   TraceOut_MoveUp[112] := BenchUut14.MoveUp;
   TraceOut_MoveLeft[112] := BenchUut14.MoveLeft;
   TraceOut_MoveRight[112] := BenchUut14.MoveRight;
   TraceOut_ActivateGrip[112] := BenchUut14.ActivateGrip;
   TraceOut_ActivateRelease[112] := BenchUut14.ActivateRelease;
   BenchCalls := BenchCalls + 1;
 113:
   BenchUut14.ManualMode := FALSE;
   BenchUut14.SingleStepMode := TRUE;
   BenchUut14.SingleCycleMode := FALSE;
   BenchUut14.ContinuousMode := FALSE;
   BenchUut14.EmergencyStop := TRUE;
   BenchUut14.Start := FALSE;
   BenchUut14.DownButton := FALSE;
   BenchUut14.UpButton := FALSE;
   BenchUut14.LeftButton := FALSE;
   BenchUut14.RightButton := FALSE;
   BenchUut14.GripButton := FALSE;
   BenchUut14.ReleaseButton := FALSE;
   BenchUut14.DownLimitSwitch := FALSE;
   BenchUut14.UpLimitSwitch := TRUE;
   BenchUut14.LeftLimitSwitch := TRUE;
   BenchUut14.RightLimitSwitch := FALSE;
   BenchUut14.GripLimitSwitch := FALSE;
   BenchUut14.ReleaseLimitSwitch := FALSE;
   TraceIn_ManualMode[113] := BenchUut14.ManualMode;
   TraceIn_SingleStepMode[113] := BenchUut14.SingleStepMode;
   TraceIn_SingleCycleMode[113] := BenchUut14.SingleCycleMode;
   TraceIn_ContinuousMode[113] := BenchUut14.ContinuousMode;
   TraceIn_EmergencyStop[113] := BenchUut14.EmergencyStop;
   TraceIn_Start[113] := BenchUut14.Start;
   TraceIn_DownButton[113] := BenchUut14.DownButton;
   TraceIn_UpButton[113] := BenchUut14.UpButton;
   TraceIn_LeftButton[113] := BenchUut14.LeftButton;
   TraceIn_RightButton[113] := BenchUut14.RightButton;
   TraceIn_GripButton[113] := BenchUut14.GripButton;
   TraceIn_ReleaseButton[113] := BenchUut14.ReleaseButton;
   TraceIn_DownLimitSwitch[113] := BenchUut14.DownLimitSwitch;
   TraceIn_UpLimitSwitch[113] := BenchUut14.UpLimitSwitch;
   TraceIn_LeftLimitSwitch[113] := BenchUut14.LeftLimitSwitch;
   TraceIn_RightLimitSwitch[113] := BenchUut14.RightLimitSwitch;
   TraceIn_GripLimitSwitch[113] := BenchUut14.GripLimitSwitch;
   TraceIn_ReleaseLimitSwitch[113] := BenchUut14.ReleaseLimitSwitch;
   BenchUut14();
   TraceOut_MoveDown[113] := BenchUut14.MoveDown;
   TraceOut_MoveUp[113] := BenchUut14.MoveUp;
   TraceOut_MoveLeft[113] := BenchUut14.MoveLeft;
   TraceOut_MoveRight[113] := BenchUut14.MoveRight;
   TraceOut_ActivateGrip[113] := BenchUut14.ActivateGrip;
   TraceOut_ActivateRelease[113] := BenchUut14.ActivateRelease;
   BenchCalls := BenchCalls + 1;
 114:
   BenchUut14.ManualMode := FALSE;
   BenchUut14.SingleStepMode := TRUE;
   BenchUut14.SingleCycleMode := FALSE;
   BenchUut14.ContinuousMode := FALSE;
   BenchUut14.EmergencyStop := TRUE;
   BenchUut14.Start := FALSE;
   BenchUut14.DownButton := FALSE;
   BenchUut14.UpButton := FALSE;
   BenchUut14.LeftButton := FALSE;
   BenchUut14.RightButton := FALSE;
   BenchUut14.GripButton := FALSE;
   BenchUut14.ReleaseButton := FALSE;
   BenchUut14.DownLimitSwitch := FALSE;
   BenchUut14.UpLimitSwitch := TRUE;
   BenchUut14.LeftLimitSwitch := TRUE;
   BenchUut14.RightLimitSwitch := FALSE;
   BenchUut14.GripLimitSwitch := FALSE;
   BenchUut14.ReleaseLimitSwitch := FALSE;
   TraceIn_ManualMode[114] := BenchUut14.ManualMode;
   TraceIn_SingleStepMode[114] := BenchUut14.SingleStepMode;
   TraceIn_SingleCycleMode[114] := BenchUut14.SingleCycleMode;
   TraceIn_ContinuousMode[114] := BenchUut14.ContinuousMode;
   TraceIn_EmergencyStop[114] := BenchUut14.EmergencyStop;
   TraceIn_Start[114] := BenchUut14.Start;
   TraceIn_DownButton[114] := BenchUut14.DownButton;
   TraceIn_UpButton[114] := BenchUut14.UpButton;
   TraceIn_LeftButton[114] := BenchUut14.LeftButton;
   TraceIn_RightButton[114] := BenchUut14.RightButton;
   TraceIn_GripButton[114] := BenchUut14.GripButton;
   TraceIn_ReleaseButton[114] := BenchUut14.ReleaseButton;
   TraceIn_DownLimitSwitch[114] := BenchUut14.DownLimitSwitch;
   TraceIn_UpLimitSwitch[114] := BenchUut14.UpLimitSwitch;
   TraceIn_LeftLimitSwitch[114] := BenchUut14.LeftLimitSwitch;
   TraceIn_RightLimitSwitch[114] := BenchUut14.RightLimitSwitch;
   TraceIn_GripLimitSwitch[114] := BenchUut14.GripLimitSwitch;
   TraceIn_ReleaseLimitSwitch[114] := BenchUut14.ReleaseLimitSwitch;
   BenchUut14();
   TraceOut_MoveDown[114] := BenchUut14.MoveDown;
   TraceOut_MoveUp[114] := BenchUut14.MoveUp;
   TraceOut_MoveLeft[114] := BenchUut14.MoveLeft;
   TraceOut_MoveRight[114] := BenchUut14.MoveRight;
   TraceOut_ActivateGrip[114] := BenchUut14.ActivateGrip;
   TraceOut_ActivateRelease[114] := BenchUut14.ActivateRelease;
   BenchCalls := BenchCalls + 1;
 115:
   BenchUut14.ManualMode := FALSE;
   BenchUut14.SingleStepMode := TRUE;
   BenchUut14.SingleCycleMode := FALSE;
   BenchUut14.ContinuousMode := FALSE;
   BenchUut14.EmergencyStop := TRUE;
   BenchUut14.Start := FALSE;
   BenchUut14.DownButton := FALSE;
   BenchUut14.UpButton := FALSE;
   BenchUut14.LeftButton := FALSE;
   BenchUut14.RightButton := FALSE;
   BenchUut14.GripButton := FALSE;
   BenchUut14.ReleaseButton := FALSE;
   BenchUut14.DownLimitSwitch := TRUE;
   BenchUut14.UpLimitSwitch := FALSE;
   BenchUut14.LeftLimitSwitch := FALSE;
   BenchUut14.RightLimitSwitch := FALSE;
   BenchUut14.GripLimitSwitch := FALSE;
   BenchUut14.ReleaseLimitSwitch := FALSE;
   TraceIn_ManualMode[115] := BenchUut14.ManualMode;
   TraceIn_SingleStepMode[115] := BenchUut14.SingleStepMode;
   TraceIn_SingleCycleMode[115] := BenchUut14.SingleCycleMode;
   TraceIn_ContinuousMode[115] := BenchUut14.ContinuousMode;
   TraceIn_EmergencyStop[115] := BenchUut14.EmergencyStop;
   TraceIn_Start[115] := BenchUut14.Start;
   TraceIn_DownButton[115] := BenchUut14.DownButton;
   TraceIn_UpButton[115] := BenchUut14.UpButton;
   TraceIn_LeftButton[115] := BenchUut14.LeftButton;
   TraceIn_RightButton[115] := BenchUut14.RightButton;
   TraceIn_GripButton[115] := BenchUut14.GripButton;
   TraceIn_ReleaseButton[115] := BenchUut14.ReleaseButton;
   TraceIn_DownLimitSwitch[115] := BenchUut14.DownLimitSwitch;
   TraceIn_UpLimitSwitch[115] := BenchUut14.UpLimitSwitch;
   TraceIn_LeftLimitSwitch[115] := BenchUut14.LeftLimitSwitch;
   TraceIn_RightLimitSwitch[115] := BenchUut14.RightLimitSwitch;
   TraceIn_GripLimitSwitch[115] := BenchUut14.GripLimitSwitch;
   TraceIn_ReleaseLimitSwitch[115] := BenchUut14.ReleaseLimitSwitch;
   BenchUut14();
   TraceOut_MoveDown[115] := BenchUut14.MoveDown;
   TraceOut_MoveUp[115] := BenchUut14.MoveUp;
   TraceOut_MoveLeft[115] := BenchUut14.MoveLeft;
   TraceOut_MoveRight[115] := BenchUut14.MoveRight;
   TraceOut_ActivateGrip[115] := BenchUut14.ActivateGrip;
   TraceOut_ActivateRelease[115] := BenchUut14.ActivateRelease;
   BenchCalls := BenchCalls + 1;
 116:
   BenchUut14.ManualMode := FALSE;
   BenchUut14.SingleStepMode := TRUE;
   BenchUut14.SingleCycleMode := FALSE;
   BenchUut14.ContinuousMode := FALSE;
   BenchUut14.EmergencyStop := TRUE;
   BenchUut14.Start := TRUE;
   BenchUut14.DownButton := FALSE;
   BenchUut14.UpButton := FALSE;
   BenchUut14.LeftButton := FALSE;
   BenchUut14.RightButton := FALSE;
   BenchUut14.GripButton := FALSE;
   BenchUut14.ReleaseButton := FALSE;
   BenchUut14.DownLimitSwitch := FALSE;
   BenchUut14.UpLimitSwitch := FALSE;
   BenchUut14.LeftLimitSwitch := FALSE;
   BenchUut14.RightLimitSwitch := FALSE;
   BenchUut14.GripLimitSwitch := FALSE;
   BenchUut14.ReleaseLimitSwitch := FALSE;
   TraceIn_ManualMode[116] := BenchUut14.ManualMode;
   TraceIn_SingleStepMode[116] := BenchUut14.SingleStepMode;
   TraceIn_SingleCycleMode[116] := BenchUut14.SingleCycleMode;
   TraceIn_ContinuousMode[116] := BenchUut14.ContinuousMode;
   TraceIn_EmergencyStop[116] := BenchUut14.EmergencyStop;
   TraceIn_Start[116] := BenchUut14.Start;
   TraceIn_DownButton[116] := BenchUut14.DownButton;
   TraceIn_UpButton[116] := BenchUut14.UpButton;
   TraceIn_LeftButton[116] := BenchUut14.LeftButton;
   TraceIn_RightButton[116] := BenchUut14.RightButton;
   TraceIn_GripButton[116] := BenchUut14.GripButton;
   TraceIn_ReleaseButton[116] := BenchUut14.ReleaseButton;
   TraceIn_DownLimitSwitch[116] := BenchUut14.DownLimitSwitch;
   TraceIn_UpLimitSwitch[116] := BenchUut14.UpLimitSwitch;
   TraceIn_LeftLimitSwitch[116] := BenchUut14.LeftLimitSwitch;
   TraceIn_RightLimitSwitch[116] := BenchUut14.RightLimitSwitch;
   TraceIn_GripLimitSwitch[116] := BenchUut14.GripLimitSwitch;
   TraceIn_ReleaseLimitSwitch[116] := BenchUut14.ReleaseLimitSwitch;
   BenchUut14();
   TraceOut_MoveDown[116] := BenchUut14.MoveDown;
   TraceOut_MoveUp[116] := BenchUut14.MoveUp;
   TraceOut_MoveLeft[116] := BenchUut14.MoveLeft;
   TraceOut_MoveRight[116] := BenchUut14.MoveRight;
   TraceOut_ActivateGrip[116] := BenchUut14.ActivateGrip;
   TraceOut_ActivateRelease[116] := BenchUut14.ActivateRelease;
   BenchCalls := BenchCalls + 1;
 117:
   BenchUut14.ManualMode := FALSE;
   BenchUut14.SingleStepMode := TRUE;
   BenchUut14.SingleCycleMode := FALSE;
   BenchUut14.ContinuousMode := FALSE;
   BenchUut14.EmergencyStop := TRUE;
   BenchUut14.Start := FALSE;
   BenchUut14.DownButton := FALSE;
   BenchUut14.UpButton := FALSE;
   BenchUut14.LeftButton := FALSE;
   BenchUut14.RightButton := FALSE;
   BenchUut14.GripButton := FALSE;
   BenchUut14.ReleaseButton := FALSE;
   BenchUut14.DownLimitSwitch := FALSE;
   BenchUut14.UpLimitSwitch := FALSE;
   BenchUut14.LeftLimitSwitch := FALSE;
   BenchUut14.RightLimitSwitch := FALSE;
   BenchUut14.GripLimitSwitch := FALSE;
   BenchUut14.ReleaseLimitSwitch := FALSE;
   TraceIn_ManualMode[117] := BenchUut14.ManualMode;
   TraceIn_SingleStepMode[117] := BenchUut14.SingleStepMode;
   TraceIn_SingleCycleMode[117] := BenchUut14.SingleCycleMode;
   TraceIn_ContinuousMode[117] := BenchUut14.ContinuousMode;
   TraceIn_EmergencyStop[117] := BenchUut14.EmergencyStop;
   TraceIn_Start[117] := BenchUut14.Start;
   TraceIn_DownButton[117] := BenchUut14.DownButton;
   TraceIn_UpButton[117] := BenchUut14.UpButton;
   TraceIn_LeftButton[117] := BenchUut14.LeftButton;
   TraceIn_RightButton[117] := BenchUut14.RightButton;
   TraceIn_GripButton[117] := BenchUut14.GripButton;
   TraceIn_ReleaseButton[117] := BenchUut14.ReleaseButton;
   TraceIn_DownLimitSwitch[117] := BenchUut14.DownLimitSwitch;
   TraceIn_UpLimitSwitch[117] := BenchUut14.UpLimitSwitch;
   TraceIn_LeftLimitSwitch[117] := BenchUut14.LeftLimitSwitch;
   TraceIn_RightLimitSwitch[117] := BenchUut14.RightLimitSwitch;
   TraceIn_GripLimitSwitch[117] := BenchUut14.GripLimitSwitch;
   TraceIn_ReleaseLimitSwitch[117] := BenchUut14.ReleaseLimitSwitch;
   BenchUut14();
   TraceOut_MoveDown[117] := BenchUut14.MoveDown;
   TraceOut_MoveUp[117] := BenchUut14.MoveUp;
   TraceOut_MoveLeft[117] := BenchUut14.MoveLeft;
   TraceOut_MoveRight[117] := BenchUut14.MoveRight;
   TraceOut_ActivateGrip[117] := BenchUut14.ActivateGrip;
   TraceOut_ActivateRelease[117] := BenchUut14.ActivateRelease;
   BenchCalls := BenchCalls + 1;
 118:
   BenchUut14.ManualMode := FALSE;
   BenchUut14.SingleStepMode := TRUE;
   BenchUut14.SingleCycleMode := FALSE;
   BenchUut14.ContinuousMode := FALSE;
   BenchUut14.EmergencyStop := TRUE;
   BenchUut14.Start := FALSE;
   BenchUut14.DownButton := FALSE;
   BenchUut14.UpButton := FALSE;
   BenchUut14.LeftButton := FALSE;
   BenchUut14.RightButton := FALSE;
   BenchUut14.GripButton := FALSE;
   BenchUut14.ReleaseButton := FALSE;
   BenchUut14.DownLimitSwitch := FALSE;
   BenchUut14.UpLimitSwitch := FALSE;
   BenchUut14.LeftLimitSwitch := FALSE;
   BenchUut14.RightLimitSwitch := FALSE;
   BenchUut14.GripLimitSwitch := FALSE;
   BenchUut14.ReleaseLimitSwitch := FALSE;
   TraceIn_ManualMode[118] := BenchUut14.ManualMode;
   TraceIn_SingleStepMode[118] := BenchUut14.SingleStepMode;
   TraceIn_SingleCycleMode[118] := BenchUut14.SingleCycleMode;
   TraceIn_ContinuousMode[118] := BenchUut14.ContinuousMode;
   TraceIn_EmergencyStop[118] := BenchUut14.EmergencyStop;
   TraceIn_Start[118] := BenchUut14.Start;
   TraceIn_DownButton[118] := BenchUut14.DownButton;
   TraceIn_UpButton[118] := BenchUut14.UpButton;
   TraceIn_LeftButton[118] := BenchUut14.LeftButton;
   TraceIn_RightButton[118] := BenchUut14.RightButton;
   TraceIn_GripButton[118] := BenchUut14.GripButton;
   TraceIn_ReleaseButton[118] := BenchUut14.ReleaseButton;
   TraceIn_DownLimitSwitch[118] := BenchUut14.DownLimitSwitch;
   TraceIn_UpLimitSwitch[118] := BenchUut14.UpLimitSwitch;
   TraceIn_LeftLimitSwitch[118] := BenchUut14.LeftLimitSwitch;
   TraceIn_RightLimitSwitch[118] := BenchUut14.RightLimitSwitch;
   TraceIn_GripLimitSwitch[118] := BenchUut14.GripLimitSwitch;
   TraceIn_ReleaseLimitSwitch[118] := BenchUut14.ReleaseLimitSwitch;
   BenchUut14();
   TraceOut_MoveDown[118] := BenchUut14.MoveDown;
   TraceOut_MoveUp[118] := BenchUut14.MoveUp;
   TraceOut_MoveLeft[118] := BenchUut14.MoveLeft;
   TraceOut_MoveRight[118] := BenchUut14.MoveRight;
   TraceOut_ActivateGrip[118] := BenchUut14.ActivateGrip;
   TraceOut_ActivateRelease[118] := BenchUut14.ActivateRelease;
   BenchCalls := BenchCalls + 1;
 119:
   BenchUut14.ManualMode := FALSE;
   BenchUut14.SingleStepMode := TRUE;
   BenchUut14.SingleCycleMode := FALSE;
   BenchUut14.ContinuousMode := FALSE;
   BenchUut14.EmergencyStop := TRUE;
   BenchUut14.Start := FALSE;
   BenchUut14.DownButton := FALSE;
   BenchUut14.UpButton := FALSE;
   BenchUut14.LeftButton := FALSE;
   BenchUut14.RightButton := FALSE;
   BenchUut14.GripButton := FALSE;
   BenchUut14.ReleaseButton := FALSE;
   BenchUut14.DownLimitSwitch := FALSE;
   BenchUut14.UpLimitSwitch := FALSE;
   BenchUut14.LeftLimitSwitch := FALSE;
   BenchUut14.RightLimitSwitch := FALSE;
   BenchUut14.GripLimitSwitch := TRUE;
   BenchUut14.ReleaseLimitSwitch := FALSE;
   TraceIn_ManualMode[119] := BenchUut14.ManualMode;
   TraceIn_SingleStepMode[119] := BenchUut14.SingleStepMode;
   TraceIn_SingleCycleMode[119] := BenchUut14.SingleCycleMode;
   TraceIn_ContinuousMode[119] := BenchUut14.ContinuousMode;
   TraceIn_EmergencyStop[119] := BenchUut14.EmergencyStop;
   TraceIn_Start[119] := BenchUut14.Start;
   TraceIn_DownButton[119] := BenchUut14.DownButton;
   TraceIn_UpButton[119] := BenchUut14.UpButton;
   TraceIn_LeftButton[119] := BenchUut14.LeftButton;
   TraceIn_RightButton[119] := BenchUut14.RightButton;
   TraceIn_GripButton[119] := BenchUut14.GripButton;
   TraceIn_ReleaseButton[119] := BenchUut14.ReleaseButton;
   TraceIn_DownLimitSwitch[119] := BenchUut14.DownLimitSwitch;
   TraceIn_UpLimitSwitch[119] := BenchUut14.UpLimitSwitch;
   TraceIn_LeftLimitSwitch[119] := BenchUut14.LeftLimitSwitch;
   TraceIn_RightLimitSwitch[119] := BenchUut14.RightLimitSwitch;
   TraceIn_GripLimitSwitch[119] := BenchUut14.GripLimitSwitch;
   TraceIn_ReleaseLimitSwitch[119] := BenchUut14.ReleaseLimitSwitch;
   BenchUut14();
   TraceOut_MoveDown[119] := BenchUut14.MoveDown;
   TraceOut_MoveUp[119] := BenchUut14.MoveUp;
   TraceOut_MoveLeft[119] := BenchUut14.MoveLeft;
   TraceOut_MoveRight[119] := BenchUut14.MoveRight;
   TraceOut_ActivateGrip[119] := BenchUut14.ActivateGrip;
   TraceOut_ActivateRelease[119] := BenchUut14.ActivateRelease;
   BenchCalls := BenchCalls + 1;
 120:
   BenchUut14.ManualMode := FALSE;
   BenchUut14.SingleStepMode := TRUE;
   BenchUut14.SingleCycleMode := FALSE;
   BenchUut14.ContinuousMode := FALSE;
   BenchUut14.EmergencyStop := TRUE;
   BenchUut14.Start := TRUE;
   BenchUut14.DownButton := FALSE;
   BenchUut14.UpButton := FALSE;
   BenchUut14.LeftButton := FALSE;
   BenchUut14.RightButton := FALSE;
   BenchUut14.GripButton := FALSE;
   BenchUut14.ReleaseButton := FALSE;
   BenchUut14.DownLimitSwitch := FALSE;
   BenchUut14.UpLimitSwitch := FALSE;
   BenchUut14.LeftLimitSwitch := FALSE;
   BenchUut14.RightLimitSwitch := FALSE;
   BenchUut14.GripLimitSwitch := FALSE;
   BenchUut14.ReleaseLimitSwitch := FALSE;
   TraceIn_ManualMode[120] := BenchUut14.ManualMode;
   TraceIn_SingleStepMode[120] := BenchUut14.SingleStepMode;
   TraceIn_SingleCycleMode[120] := BenchUut14.SingleCycleMode;
   TraceIn_ContinuousMode[120] := BenchUut14.ContinuousMode;
   TraceIn_EmergencyStop[120] := BenchUut14.EmergencyStop;
   TraceIn_Start[120] := BenchUut14.Start;
   TraceIn_DownButton[120] := BenchUut14.DownButton;
   TraceIn_UpButton[120] := BenchUut14.UpButton;
   TraceIn_LeftButton[120] := BenchUut14.LeftButton;
   TraceIn_RightButton[120] := BenchUut14.RightButton;
   TraceIn_GripButton[120] := BenchUut14.GripButton;
   TraceIn_ReleaseButton[120] := BenchUut14.ReleaseButton;
   TraceIn_DownLimitSwitch[120] := BenchUut14.DownLimitSwitch;
   TraceIn_UpLimitSwitch[120] := BenchUut14.UpLimitSwitch;
   TraceIn_LeftLimitSwitch[120] := BenchUut14.LeftLimitSwitch;
   TraceIn_RightLimitSwitch[120] := BenchUut14.RightLimitSwitch;
   TraceIn_GripLimitSwitch[120] := BenchUut14.GripLimitSwitch;
   TraceIn_ReleaseLimitSwitch[120] := BenchUut14.ReleaseLimitSwitch;
   BenchUut14();
   TraceOut_MoveDown[120] := BenchUut14.MoveDown;
   TraceOut_MoveUp[120] := BenchUut14.MoveUp;
   TraceOut_MoveLeft[120] := BenchUut14.MoveLeft;
   TraceOut_MoveRight[120] := BenchUut14.MoveRight;
   TraceOut_ActivateGrip[120] := BenchUut14.ActivateGrip;
   TraceOut_ActivateRelease[120] := BenchUut14.ActivateRelease;
   BenchCalls := BenchCalls + 1;
 121:
   BenchUut14.ManualMode := FALSE;
   BenchUut14.SingleStepMode := TRUE;
   BenchUut14.SingleCycleMode := FALSE;
   BenchUut14.ContinuousMode := FALSE;
   BenchUut14.EmergencyStop := TRUE;
   BenchUut14.Start := FALSE;
   BenchUut14.DownButton := FALSE;
   BenchUut14.UpButton := FALSE;
   BenchUut14.LeftButton := FALSE;
   BenchUut14.RightButton := FALSE;
   BenchUut14.GripButton := FALSE;
   BenchUut14.ReleaseButton := FALSE;
   BenchUut14.DownLimitSwitch := FALSE;
   BenchUut14.UpLimitSwitch := FALSE;
   BenchUut14.LeftLimitSwitch := FALSE;
   BenchUut14.RightLimitSwitch := FALSE;
   BenchUut14.GripLimitSwitch := FALSE;
   BenchUut14.ReleaseLimitSwitch := FALSE;
   TraceIn_ManualMode[121] := BenchUut14.ManualMode;
   TraceIn_SingleStepMode[121] := BenchUut14.SingleStepMode;
   TraceIn_SingleCycleMode[121] := BenchUut14.SingleCycleMode;
   TraceIn_ContinuousMode[121] := BenchUut14.ContinuousMode;
   TraceIn_EmergencyStop[121] := BenchUut14.EmergencyStop;
   TraceIn_Start[121] := BenchUut14.Start;
   TraceIn_DownButton[121] := BenchUut14.DownButton;
   TraceIn_UpButton[121] := BenchUut14.UpButton;
   TraceIn_LeftButton[121] := BenchUut14.LeftButton;
   TraceIn_RightButton[121] := BenchUut14.RightButton;
   TraceIn_GripButton[121] := BenchUut14.GripButton;
   TraceIn_ReleaseButton[121] := BenchUut14.ReleaseButton;
   TraceIn_DownLimitSwitch[121] := BenchUut14.DownLimitSwitch;
   TraceIn_UpLimitSwitch[121] := BenchUut14.UpLimitSwitch;
   TraceIn_LeftLimitSwitch[121] := BenchUut14.LeftLimitSwitch;
   TraceIn_RightLimitSwitch[121] := BenchUut14.RightLimitSwitch;
   TraceIn_GripLimitSwitch[121] := BenchUut14.GripLimitSwitch;
   TraceIn_ReleaseLimitSwitch[121] := BenchUut14.ReleaseLimitSwitch;
   BenchUut14();
   TraceOut_MoveDown[121] := BenchUut14.MoveDown;
   TraceOut_MoveUp[121] := BenchUut14.MoveUp;
   TraceOut_MoveLeft[121] := BenchUut14.MoveLeft;
   TraceOut_MoveRight[121] := BenchUut14.MoveRight;
   TraceOut_ActivateGrip[121] := BenchUut14.ActivateGrip;
   TraceOut_ActivateRelease[121] := BenchUut14.ActivateRelease;
   BenchCalls := BenchCalls + 1;
 122:
   BenchUut14.ManualMode := FALSE;
   BenchUut14.SingleStepMode := TRUE;
   BenchUut14.SingleCycleMode := FALSE;
   BenchUut14.ContinuousMode := FALSE;
   BenchUut14.EmergencyStop := TRUE;
   BenchUut14.Start := FALSE;
   BenchUut14.DownButton := FALSE;
   BenchUut14.UpButton := FALSE;
   BenchUut14.LeftButton := FALSE;
   BenchUut14.RightButton := FALSE;
   BenchUut14.GripButton := FALSE;
   BenchUut14.ReleaseButton := FALSE;
   BenchUut14.DownLimitSwitch := FALSE;
   BenchUut14.UpLimitSwitch := FALSE;
   BenchUut14.LeftLimitSwitch := FALSE;
   BenchUut14.RightLimitSwitch := FALSE;
   BenchUut14.GripLimitSwitch := FALSE;
   BenchUut14.ReleaseLimitSwitch := FALSE;
   TraceIn_ManualMode[122] := BenchUut14.ManualMode;
   TraceIn_SingleStepMode[122] := BenchUut14.SingleStepMode;
   TraceIn_SingleCycleMode[122] := BenchUut14.SingleCycleMode;
   TraceIn_ContinuousMode[122] := BenchUut14.ContinuousMode;
   TraceIn_EmergencyStop[122] := BenchUut14.EmergencyStop;
   TraceIn_Start[122] := BenchUut14.Start;
   TraceIn_DownButton[122] := BenchUut14.DownButton;
   TraceIn_UpButton[122] := BenchUut14.UpButton;
   TraceIn_LeftButton[122] := BenchUut14.LeftButton;
   TraceIn_RightButton[122] := BenchUut14.RightButton;
   TraceIn_GripButton[122] := BenchUut14.GripButton;
   TraceIn_ReleaseButton[122] := BenchUut14.ReleaseButton;
   TraceIn_DownLimitSwitch[122] := BenchUut14.DownLimitSwitch;
   TraceIn_UpLimitSwitch[122] := BenchUut14.UpLimitSwitch;
   TraceIn_LeftLimitSwitch[122] := BenchUut14.LeftLimitSwitch;
   TraceIn_RightLimitSwitch[122] := BenchUut14.RightLimitSwitch;
   TraceIn_GripLimitSwitch[122] := BenchUut14.GripLimitSwitch;
   TraceIn_ReleaseLimitSwitch[122] := BenchUut14.ReleaseLimitSwitch;
   BenchUut14();
   TraceOut_MoveDown[122] := BenchUut14.MoveDown;
   TraceOut_MoveUp[122] := BenchUut14.MoveUp;
   TraceOut_MoveLeft[122] := BenchUut14.MoveLeft;
   TraceOut_MoveRight[122] := BenchUut14.MoveRight;
   TraceOut_ActivateGrip[122] := BenchUut14.ActivateGrip;
   TraceOut_ActivateRelease[122] := BenchUut14.ActivateRelease;
   BenchCalls := BenchCalls + 1;
 123:
   BenchUut14.ManualMode := FALSE;
   BenchUut14.SingleStepMode := TRUE;
   BenchUut14.SingleCycleMode := FALSE;
   BenchUut14.ContinuousMode := FALSE;
   BenchUut14.EmergencyStop := TRUE;
   BenchUut14.Start := FALSE;
   BenchUut14.DownButton := FALSE;
   BenchUut14.UpButton := FALSE;
   BenchUut14.LeftButton := FALSE;
   BenchUut14.RightButton := FALSE;
   BenchUut14.GripButton := FALSE;
   BenchUut14.ReleaseButton := FALSE;
   BenchUut14.DownLimitSwitch := FALSE;
   BenchUut14.UpLimitSwitch := TRUE;
   BenchUut14.LeftLimitSwitch := FALSE;
   BenchUut14.RightLimitSwitch := FALSE;
   BenchUut14.GripLimitSwitch := FALSE;
   BenchUut14.ReleaseLimitSwitch := FALSE;
   TraceIn_ManualMode[123] := BenchUut14.ManualMode;
   TraceIn_SingleStepMode[123] := BenchUut14.SingleStepMode;
   TraceIn_SingleCycleMode[123] := BenchUut14.SingleCycleMode;
   TraceIn_ContinuousMode[123] := BenchUut14.ContinuousMode;
   TraceIn_EmergencyStop[123] := BenchUut14.EmergencyStop;
   TraceIn_Start[123] := BenchUut14.Start;
   TraceIn_DownButton[123] := BenchUut14.DownButton;
   TraceIn_UpButton[123] := BenchUut14.UpButton;
   TraceIn_LeftButton[123] := BenchUut14.LeftButton;
   TraceIn_RightButton[123] := BenchUut14.RightButton;
   TraceIn_GripButton[123] := BenchUut14.GripButton;
   TraceIn_ReleaseButton[123] := BenchUut14.ReleaseButton;
   TraceIn_DownLimitSwitch[123] := BenchUut14.DownLimitSwitch;
   TraceIn_UpLimitSwitch[123] := BenchUut14.UpLimitSwitch;
   TraceIn_LeftLimitSwitch[123] := BenchUut14.LeftLimitSwitch;
   TraceIn_RightLimitSwitch[123] := BenchUut14.RightLimitSwitch;
   TraceIn_GripLimitSwitch[123] := BenchUut14.GripLimitSwitch;
   TraceIn_ReleaseLimitSwitch[123] := BenchUut14.ReleaseLimitSwitch;
   BenchUut14();
   TraceOut_MoveDown[123] := BenchUut14.MoveDown;
   TraceOut_MoveUp[123] := BenchUut14.MoveUp;
   TraceOut_MoveLeft[123] := BenchUut14.MoveLeft;
   TraceOut_MoveRight[123] := BenchUut14.MoveRight;
   TraceOut_ActivateGrip[123] := BenchUut14.ActivateGrip;
   TraceOut_ActivateRelease[123] := BenchUut14.ActivateRelease;
   BenchCalls := BenchCalls + 1;
 124:
   BenchUut14.ManualMode := FALSE;
   BenchUut14.SingleStepMode := TRUE;
   BenchUut14.SingleCycleMode := FALSE;
   BenchUut14.ContinuousMode := FALSE;
   BenchUut14.EmergencyStop := TRUE;
   BenchUut14.Start := TRUE;
   BenchUut14.DownButton := FALSE;
   BenchUut14.UpButton := FALSE;
   BenchUut14.LeftButton := FALSE;
   BenchUut14.RightButton := FALSE;
   BenchUut14.GripButton := FALSE;
   BenchUut14.ReleaseButton := FALSE;
   BenchUut14.DownLimitSwitch := FALSE;
   BenchUut14.UpLimitSwitch := FALSE;
   BenchUut14.LeftLimitSwitch := FALSE;
   BenchUut14.RightLimitSwitch := FALSE;
   BenchUut14.GripLimitSwitch := FALSE;
   BenchUut14.ReleaseLimitSwitch := FALSE;
   TraceIn_ManualMode[124] := BenchUut14.ManualMode;
   TraceIn_SingleStepMode[124] := BenchUut14.SingleStepMode;
   TraceIn_SingleCycleMode[124] := BenchUut14.SingleCycleMode;
   TraceIn_ContinuousMode[124] := BenchUut14.ContinuousMode;
   TraceIn_EmergencyStop[124] := BenchUut14.EmergencyStop;
   TraceIn_Start[124] := BenchUut14.Start;
   TraceIn_DownButton[124] := BenchUut14.DownButton;
   TraceIn_UpButton[124] := BenchUut14.UpButton;
   TraceIn_LeftButton[124] := BenchUut14.LeftButton;
   TraceIn_RightButton[124] := BenchUut14.RightButton;
   TraceIn_GripButton[124] := BenchUut14.GripButton;
   TraceIn_ReleaseButton[124] := BenchUut14.ReleaseButton;
   TraceIn_DownLimitSwitch[124] := BenchUut14.DownLimitSwitch;
   TraceIn_UpLimitSwitch[124] := BenchUut14.UpLimitSwitch;
   TraceIn_LeftLimitSwitch[124] := BenchUut14.LeftLimitSwitch;
   TraceIn_RightLimitSwitch[124] := BenchUut14.RightLimitSwitch;
   TraceIn_GripLimitSwitch[124] := BenchUut14.GripLimitSwitch;
   TraceIn_ReleaseLimitSwitch[124] := BenchUut14.ReleaseLimitSwitch;
   BenchUut14();
   TraceOut_MoveDown[124] := BenchUut14.MoveDown;
   TraceOut_MoveUp[124] := BenchUut14.MoveUp;
   TraceOut_MoveLeft[124] := BenchUut14.MoveLeft;
   TraceOut_MoveRight[124] := BenchUut14.MoveRight;
   TraceOut_ActivateGrip[124] := BenchUut14.ActivateGrip;
   TraceOut_ActivateRelease[124] := BenchUut14.ActivateRelease;
   BenchCalls := BenchCalls + 1;
 125:
   BenchUut14.ManualMode := FALSE;
   BenchUut14.SingleStepMode := TRUE;
   BenchUut14.SingleCycleMode := FALSE;
   BenchUut14.ContinuousMode := FALSE;
   BenchUut14.EmergencyStop := TRUE;
   BenchUut14.Start := FALSE;
   BenchUut14.DownButton := FALSE;
   BenchUut14.UpButton := FALSE;
   BenchUut14.LeftButton := FALSE;
   BenchUut14.RightButton := FALSE;
   BenchUut14.GripButton := FALSE;
   BenchUut14.ReleaseButton := FALSE;
   BenchUut14.DownLimitSwitch := FALSE;
   BenchUut14.UpLimitSwitch := FALSE;
   BenchUut14.LeftLimitSwitch := FALSE;
   BenchUut14.RightLimitSwitch := FALSE;
   BenchUut14.GripLimitSwitch := FALSE;
   BenchUut14.ReleaseLimitSwitch := FALSE;
   TraceIn_ManualMode[125] := BenchUut14.ManualMode;
   TraceIn_SingleStepMode[125] := BenchUut14.SingleStepMode;
   TraceIn_SingleCycleMode[125] := BenchUut14.SingleCycleMode;
   TraceIn_ContinuousMode[125] := BenchUut14.ContinuousMode;
   TraceIn_EmergencyStop[125] := BenchUut14.EmergencyStop;
   TraceIn_Start[125] := BenchUut14.Start;
   TraceIn_DownButton[125] := BenchUut14.DownButton;
   TraceIn_UpButton[125] := BenchUut14.UpButton;
   TraceIn_LeftButton[125] := BenchUut14.LeftButton;
   TraceIn_RightButton[125] := BenchUut14.RightButton;
   TraceIn_GripButton[125] := BenchUut14.GripButton;
   TraceIn_ReleaseButton[125] := BenchUut14.ReleaseButton;
   TraceIn_DownLimitSwitch[125] := BenchUut14.DownLimitSwitch;
   TraceIn_UpLimitSwitch[125] := BenchUut14.UpLimitSwitch;
   TraceIn_LeftLimitSwitch[125] := BenchUut14.LeftLimitSwitch;
   TraceIn_RightLimitSwitch[125] := BenchUut14.RightLimitSwitch;
   TraceIn_GripLimitSwitch[125] := BenchUut14.GripLimitSwitch;
   TraceIn_ReleaseLimitSwitch[125] := BenchUut14.ReleaseLimitSwitch;
   BenchUut14();
   TraceOut_MoveDown[125] := BenchUut14.MoveDown;
   TraceOut_MoveUp[125] := BenchUut14.MoveUp;
   TraceOut_MoveLeft[125] := BenchUut14.MoveLeft;
   TraceOut_MoveRight[125] := BenchUut14.MoveRight;
   TraceOut_ActivateGrip[125] := BenchUut14.ActivateGrip;
   TraceOut_ActivateRelease[125] := BenchUut14.ActivateRelease;
   BenchCalls := BenchCalls + 1;
 126:
   BenchUut14.ManualMode := FALSE;
   BenchUut14.SingleStepMode := TRUE;
   BenchUut14.SingleCycleMode := FALSE;
   BenchUut14.ContinuousMode := FALSE;
   BenchUut14.EmergencyStop := TRUE;
   BenchUut14.Start := FALSE;
   BenchUut14.DownButton := FALSE;
   BenchUut14.UpButton := FALSE;
   BenchUut14.LeftButton := FALSE;
   BenchUut14.RightButton := FALSE;
   BenchUut14.GripButton := FALSE;
   BenchUut14.ReleaseButton := FALSE;
   BenchUut14.DownLimitSwitch := FALSE;
   BenchUut14.UpLimitSwitch := FALSE;
   BenchUut14.LeftLimitSwitch := FALSE;
   BenchUut14.RightLimitSwitch := FALSE;
   BenchUut14.GripLimitSwitch := FALSE;
   BenchUut14.ReleaseLimitSwitch := FALSE;
   TraceIn_ManualMode[126] := BenchUut14.ManualMode;
   TraceIn_SingleStepMode[126] := BenchUut14.SingleStepMode;
   TraceIn_SingleCycleMode[126] := BenchUut14.SingleCycleMode;
   TraceIn_ContinuousMode[126] := BenchUut14.ContinuousMode;
   TraceIn_EmergencyStop[126] := BenchUut14.EmergencyStop;
   TraceIn_Start[126] := BenchUut14.Start;
   TraceIn_DownButton[126] := BenchUut14.DownButton;
   TraceIn_UpButton[126] := BenchUut14.UpButton;
   TraceIn_LeftButton[126] := BenchUut14.LeftButton;
   TraceIn_RightButton[126] := BenchUut14.RightButton;
   TraceIn_GripButton[126] := BenchUut14.GripButton;
   TraceIn_ReleaseButton[126] := BenchUut14.ReleaseButton;
   TraceIn_DownLimitSwitch[126] := BenchUut14.DownLimitSwitch;
   TraceIn_UpLimitSwitch[126] := BenchUut14.UpLimitSwitch;
   TraceIn_LeftLimitSwitch[126] := BenchUut14.LeftLimitSwitch;
   TraceIn_RightLimitSwitch[126] := BenchUut14.RightLimitSwitch;
   TraceIn_GripLimitSwitch[126] := BenchUut14.GripLimitSwitch;
   TraceIn_ReleaseLimitSwitch[126] := BenchUut14.ReleaseLimitSwitch;
   BenchUut14();
   TraceOut_MoveDown[126] := BenchUut14.MoveDown;
   TraceOut_MoveUp[126] := BenchUut14.MoveUp;
   TraceOut_MoveLeft[126] := BenchUut14.MoveLeft;
   TraceOut_MoveRight[126] := BenchUut14.MoveRight;
   TraceOut_ActivateGrip[126] := BenchUut14.ActivateGrip;
   TraceOut_ActivateRelease[126] := BenchUut14.ActivateRelease;
   BenchCalls := BenchCalls + 1;
 127:
   BenchUut14.ManualMode := FALSE;
   BenchUut14.SingleStepMode := TRUE;
   BenchUut14.SingleCycleMode := FALSE;
   BenchUut14.ContinuousMode := FALSE;
   BenchUut14.EmergencyStop := TRUE;
   BenchUut14.Start := FALSE;
   BenchUut14.DownButton := FALSE;
   BenchUut14.UpButton := FALSE;
   BenchUut14.LeftButton := FALSE;
   BenchUut14.RightButton := FALSE;
   BenchUut14.GripButton := FALSE;
   BenchUut14.ReleaseButton := FALSE;
   BenchUut14.DownLimitSwitch := FALSE;
   BenchUut14.UpLimitSwitch := FALSE;
   BenchUut14.LeftLimitSwitch := FALSE;
   BenchUut14.RightLimitSwitch := TRUE;
   BenchUut14.GripLimitSwitch := FALSE;
   BenchUut14.ReleaseLimitSwitch := FALSE;
   TraceIn_ManualMode[127] := BenchUut14.ManualMode;
   TraceIn_SingleStepMode[127] := BenchUut14.SingleStepMode;
   TraceIn_SingleCycleMode[127] := BenchUut14.SingleCycleMode;
   TraceIn_ContinuousMode[127] := BenchUut14.ContinuousMode;
   TraceIn_EmergencyStop[127] := BenchUut14.EmergencyStop;
   TraceIn_Start[127] := BenchUut14.Start;
   TraceIn_DownButton[127] := BenchUut14.DownButton;
   TraceIn_UpButton[127] := BenchUut14.UpButton;
   TraceIn_LeftButton[127] := BenchUut14.LeftButton;
   TraceIn_RightButton[127] := BenchUut14.RightButton;
   TraceIn_GripButton[127] := BenchUut14.GripButton;
   TraceIn_ReleaseButton[127] := BenchUut14.ReleaseButton;
   TraceIn_DownLimitSwitch[127] := BenchUut14.DownLimitSwitch;
   TraceIn_UpLimitSwitch[127] := BenchUut14.UpLimitSwitch;
   TraceIn_LeftLimitSwitch[127] := BenchUut14.LeftLimitSwitch;
   TraceIn_RightLimitSwitch[127] := BenchUut14.RightLimitSwitch;
   TraceIn_GripLimitSwitch[127] := BenchUut14.GripLimitSwitch;
   TraceIn_ReleaseLimitSwitch[127] := BenchUut14.ReleaseLimitSwitch;
   BenchUut14();
   TraceOut_MoveDown[127] := BenchUut14.MoveDown;
   TraceOut_MoveUp[127] := BenchUut14.MoveUp;
   TraceOut_MoveLeft[127] := BenchUut14.MoveLeft;
   TraceOut_MoveRight[127] := BenchUut14.MoveRight;
   TraceOut_ActivateGrip[127] := BenchUut14.ActivateGrip;
   TraceOut_ActivateRelease[127] := BenchUut14.ActivateRelease;
   BenchCalls := BenchCalls + 1;
 128:
   BenchUut14.ManualMode := FALSE;
   BenchUut14.SingleStepMode := TRUE;
   BenchUut14.SingleCycleMode := FALSE;
   BenchUut14.ContinuousMode := FALSE;
   BenchUut14.EmergencyStop := TRUE;
   BenchUut14.Start := TRUE;
   BenchUut14.DownButton := FALSE;
   BenchUut14.UpButton := FALSE;
   BenchUut14.LeftButton := FALSE;
   BenchUut14.RightButton := FALSE;
   BenchUut14.GripButton := FALSE;
   BenchUut14.ReleaseButton := FALSE;
   BenchUut14.DownLimitSwitch := FALSE;
   BenchUut14.UpLimitSwitch := FALSE;
   BenchUut14.LeftLimitSwitch := FALSE;
   BenchUut14.RightLimitSwitch := FALSE;
   BenchUut14.GripLimitSwitch := FALSE;
   BenchUut14.ReleaseLimitSwitch := FALSE;
   TraceIn_ManualMode[128] := BenchUut14.ManualMode;
   TraceIn_SingleStepMode[128] := BenchUut14.SingleStepMode;
   TraceIn_SingleCycleMode[128] := BenchUut14.SingleCycleMode;
   TraceIn_ContinuousMode[128] := BenchUut14.ContinuousMode;
   TraceIn_EmergencyStop[128] := BenchUut14.EmergencyStop;
   TraceIn_Start[128] := BenchUut14.Start;
   TraceIn_DownButton[128] := BenchUut14.DownButton;
   TraceIn_UpButton[128] := BenchUut14.UpButton;
   TraceIn_LeftButton[128] := BenchUut14.LeftButton;
   TraceIn_RightButton[128] := BenchUut14.RightButton;
   TraceIn_GripButton[128] := BenchUut14.GripButton;
   TraceIn_ReleaseButton[128] := BenchUut14.ReleaseButton;
   TraceIn_DownLimitSwitch[128] := BenchUut14.DownLimitSwitch;
   TraceIn_UpLimitSwitch[128] := BenchUut14.UpLimitSwitch;
   TraceIn_LeftLimitSwitch[128] := BenchUut14.LeftLimitSwitch;
   TraceIn_RightLimitSwitch[128] := BenchUut14.RightLimitSwitch;
   TraceIn_GripLimitSwitch[128] := BenchUut14.GripLimitSwitch;
   TraceIn_ReleaseLimitSwitch[128] := BenchUut14.ReleaseLimitSwitch;
   BenchUut14();
   TraceOut_MoveDown[128] := BenchUut14.MoveDown;
   TraceOut_MoveUp[128] := BenchUut14.MoveUp;
   TraceOut_MoveLeft[128] := BenchUut14.MoveLeft;
   TraceOut_MoveRight[128] := BenchUut14.MoveRight;
   TraceOut_ActivateGrip[128] := BenchUut14.ActivateGrip;
   TraceOut_ActivateRelease[128] := BenchUut14.ActivateRelease;
   BenchCalls := BenchCalls + 1;
 129:
   BenchUut14.ManualMode := FALSE;
   BenchUut14.SingleStepMode := TRUE;
   BenchUut14.SingleCycleMode := FALSE;
   BenchUut14.ContinuousMode := FALSE;
   BenchUut14.EmergencyStop := TRUE;
   BenchUut14.Start := FALSE;
   BenchUut14.DownButton := FALSE;
   BenchUut14.UpButton := FALSE;
   BenchUut14.LeftButton := FALSE;
   BenchUut14.RightButton := FALSE;
   BenchUut14.GripButton := FALSE;
   BenchUut14.ReleaseButton := FALSE;
   BenchUut14.DownLimitSwitch := FALSE;
   BenchUut14.UpLimitSwitch := FALSE;
   BenchUut14.LeftLimitSwitch := FALSE;
   BenchUut14.RightLimitSwitch := FALSE;
   BenchUut14.GripLimitSwitch := FALSE;
   BenchUut14.ReleaseLimitSwitch := FALSE;
   TraceIn_ManualMode[129] := BenchUut14.ManualMode;
   TraceIn_SingleStepMode[129] := BenchUut14.SingleStepMode;
   TraceIn_SingleCycleMode[129] := BenchUut14.SingleCycleMode;
   TraceIn_ContinuousMode[129] := BenchUut14.ContinuousMode;
   TraceIn_EmergencyStop[129] := BenchUut14.EmergencyStop;
   TraceIn_Start[129] := BenchUut14.Start;
   TraceIn_DownButton[129] := BenchUut14.DownButton;
   TraceIn_UpButton[129] := BenchUut14.UpButton;
   TraceIn_LeftButton[129] := BenchUut14.LeftButton;
   TraceIn_RightButton[129] := BenchUut14.RightButton;
   TraceIn_GripButton[129] := BenchUut14.GripButton;
   TraceIn_ReleaseButton[129] := BenchUut14.ReleaseButton;
   TraceIn_DownLimitSwitch[129] := BenchUut14.DownLimitSwitch;
   TraceIn_UpLimitSwitch[129] := BenchUut14.UpLimitSwitch;
   TraceIn_LeftLimitSwitch[129] := BenchUut14.LeftLimitSwitch;
   TraceIn_RightLimitSwitch[129] := BenchUut14.RightLimitSwitch;
   TraceIn_GripLimitSwitch[129] := BenchUut14.GripLimitSwitch;
   TraceIn_ReleaseLimitSwitch[129] := BenchUut14.ReleaseLimitSwitch;
   BenchUut14();
   TraceOut_MoveDown[129] := BenchUut14.MoveDown;
   TraceOut_MoveUp[129] := BenchUut14.MoveUp;
   TraceOut_MoveLeft[129] := BenchUut14.MoveLeft;
   TraceOut_MoveRight[129] := BenchUut14.MoveRight;
   TraceOut_ActivateGrip[129] := BenchUut14.ActivateGrip;
   TraceOut_ActivateRelease[129] := BenchUut14.ActivateRelease;
   BenchCalls := BenchCalls + 1;
 130:
   BenchUut14.ManualMode := FALSE;
   BenchUut14.SingleStepMode := TRUE;
   BenchUut14.SingleCycleMode := FALSE;
   BenchUut14.ContinuousMode := FALSE;
   BenchUut14.EmergencyStop := TRUE;
   BenchUut14.Start := FALSE;
   BenchUut14.DownButton := FALSE;
   BenchUut14.UpButton := FALSE;
   BenchUut14.LeftButton := FALSE;
   BenchUut14.RightButton := FALSE;
   BenchUut14.GripButton := FALSE;
   BenchUut14.ReleaseButton := FALSE;
   BenchUut14.DownLimitSwitch := FALSE;
   BenchUut14.UpLimitSwitch := FALSE;
   BenchUut14.LeftLimitSwitch := FALSE;
   BenchUut14.RightLimitSwitch := FALSE;
   BenchUut14.GripLimitSwitch := FALSE;
   BenchUut14.ReleaseLimitSwitch := FALSE;
   TraceIn_ManualMode[130] := BenchUut14.ManualMode;
   TraceIn_SingleStepMode[130] := BenchUut14.SingleStepMode;
   TraceIn_SingleCycleMode[130] := BenchUut14.SingleCycleMode;
   TraceIn_ContinuousMode[130] := BenchUut14.ContinuousMode;
   TraceIn_EmergencyStop[130] := BenchUut14.EmergencyStop;
   TraceIn_Start[130] := BenchUut14.Start;
   TraceIn_DownButton[130] := BenchUut14.DownButton;
   TraceIn_UpButton[130] := BenchUut14.UpButton;
   TraceIn_LeftButton[130] := BenchUut14.LeftButton;
   TraceIn_RightButton[130] := BenchUut14.RightButton;
   TraceIn_GripButton[130] := BenchUut14.GripButton;
   TraceIn_ReleaseButton[130] := BenchUut14.ReleaseButton;
   TraceIn_DownLimitSwitch[130] := BenchUut14.DownLimitSwitch;
   TraceIn_UpLimitSwitch[130] := BenchUut14.UpLimitSwitch;
   TraceIn_LeftLimitSwitch[130] := BenchUut14.LeftLimitSwitch;
   TraceIn_RightLimitSwitch[130] := BenchUut14.RightLimitSwitch;
   TraceIn_GripLimitSwitch[130] := BenchUut14.GripLimitSwitch;
   TraceIn_ReleaseLimitSwitch[130] := BenchUut14.ReleaseLimitSwitch;
   BenchUut14();
   TraceOut_MoveDown[130] := BenchUut14.MoveDown;
   TraceOut_MoveUp[130] := BenchUut14.MoveUp;
   TraceOut_MoveLeft[130] := BenchUut14.MoveLeft;
   TraceOut_MoveRight[130] := BenchUut14.MoveRight;
   TraceOut_ActivateGrip[130] := BenchUut14.ActivateGrip;
   TraceOut_ActivateRelease[130] := BenchUut14.ActivateRelease;
   BenchCalls := BenchCalls + 1;
 131:
   BenchUut14.ManualMode := FALSE;
   BenchUut14.SingleStepMode := TRUE;
   BenchUut14.SingleCycleMode := FALSE;
   BenchUut14.ContinuousMode := FALSE;
   BenchUut14.EmergencyStop := TRUE;
   BenchUut14.Start := FALSE;
   BenchUut14.DownButton := FALSE;
   BenchUut14.UpButton := FALSE;
   BenchUut14.LeftButton := FALSE;
   BenchUut14.RightButton := FALSE;
   BenchUut14.GripButton := FALSE;
   BenchUut14.ReleaseButton := FALSE;
   BenchUut14.DownLimitSwitch := TRUE;
   BenchUut14.UpLimitSwitch := FALSE;
   BenchUut14.LeftLimitSwitch := FALSE;
   BenchUut14.RightLimitSwitch := FALSE;
   BenchUut14.GripLimitSwitch := FALSE;
   BenchUut14.ReleaseLimitSwitch := FALSE;
   TraceIn_ManualMode[131] := BenchUut14.ManualMode;
   TraceIn_SingleStepMode[131] := BenchUut14.SingleStepMode;
   TraceIn_SingleCycleMode[131] := BenchUut14.SingleCycleMode;
   TraceIn_ContinuousMode[131] := BenchUut14.ContinuousMode;
   TraceIn_EmergencyStop[131] := BenchUut14.EmergencyStop;
   TraceIn_Start[131] := BenchUut14.Start;
   TraceIn_DownButton[131] := BenchUut14.DownButton;
   TraceIn_UpButton[131] := BenchUut14.UpButton;
   TraceIn_LeftButton[131] := BenchUut14.LeftButton;
   TraceIn_RightButton[131] := BenchUut14.RightButton;
   TraceIn_GripButton[131] := BenchUut14.GripButton;
   TraceIn_ReleaseButton[131] := BenchUut14.ReleaseButton;
   TraceIn_DownLimitSwitch[131] := BenchUut14.DownLimitSwitch;
   TraceIn_UpLimitSwitch[131] := BenchUut14.UpLimitSwitch;
   TraceIn_LeftLimitSwitch[131] := BenchUut14.LeftLimitSwitch;
   TraceIn_RightLimitSwitch[131] := BenchUut14.RightLimitSwitch;
   TraceIn_GripLimitSwitch[131] := BenchUut14.GripLimitSwitch;
   TraceIn_ReleaseLimitSwitch[131] := BenchUut14.ReleaseLimitSwitch;
   BenchUut14();
   TraceOut_MoveDown[131] := BenchUut14.MoveDown;
   TraceOut_MoveUp[131] := BenchUut14.MoveUp;
   TraceOut_MoveLeft[131] := BenchUut14.MoveLeft;
   TraceOut_MoveRight[131] := BenchUut14.MoveRight;
   TraceOut_ActivateGrip[131] := BenchUut14.ActivateGrip;
   TraceOut_ActivateRelease[131] := BenchUut14.ActivateRelease;
   BenchCalls := BenchCalls + 1;
 132:
   BenchUut14.ManualMode := FALSE;
   BenchUut14.SingleStepMode := TRUE;
   BenchUut14.SingleCycleMode := FALSE;
   BenchUut14.ContinuousMode := FALSE;
   BenchUut14.EmergencyStop := TRUE;
   BenchUut14.Start := TRUE;
   BenchUut14.DownButton := FALSE;
   BenchUut14.UpButton := FALSE;
   BenchUut14.LeftButton := FALSE;
   BenchUut14.RightButton := FALSE;
   BenchUut14.GripButton := FALSE;
   BenchUut14.ReleaseButton := FALSE;
   BenchUut14.DownLimitSwitch := FALSE;
   BenchUut14.UpLimitSwitch := FALSE;
   BenchUut14.LeftLimitSwitch := FALSE;
   BenchUut14.RightLimitSwitch := FALSE;
   BenchUut14.GripLimitSwitch := FALSE;
   BenchUut14.ReleaseLimitSwitch := FALSE;
   TraceIn_ManualMode[132] := BenchUut14.ManualMode;
   TraceIn_SingleStepMode[132] := BenchUut14.SingleStepMode;
   TraceIn_SingleCycleMode[132] := BenchUut14.SingleCycleMode;
   TraceIn_ContinuousMode[132] := BenchUut14.ContinuousMode;
   TraceIn_EmergencyStop[132] := BenchUut14.EmergencyStop;
   TraceIn_Start[132] := BenchUut14.Start;
   TraceIn_DownButton[132] := BenchUut14.DownButton;
   TraceIn_UpButton[132] := BenchUut14.UpButton;
   TraceIn_LeftButton[132] := BenchUut14.LeftButton;
   TraceIn_RightButton[132] := BenchUut14.RightButton;
   TraceIn_GripButton[132] := BenchUut14.GripButton;
   TraceIn_ReleaseButton[132] := BenchUut14.ReleaseButton;
   TraceIn_DownLimitSwitch[132] := BenchUut14.DownLimitSwitch;
   TraceIn_UpLimitSwitch[132] := BenchUut14.UpLimitSwitch;
   TraceIn_LeftLimitSwitch[132] := BenchUut14.LeftLimitSwitch;
   TraceIn_RightLimitSwitch[132] := BenchUut14.RightLimitSwitch;
   TraceIn_GripLimitSwitch[132] := BenchUut14.GripLimitSwitch;
   TraceIn_ReleaseLimitSwitch[132] := BenchUut14.ReleaseLimitSwitch;
   BenchUut14();
   TraceOut_MoveDown[132] := BenchUut14.MoveDown;
   TraceOut_MoveUp[132] := BenchUut14.MoveUp;
   TraceOut_MoveLeft[132] := BenchUut14.MoveLeft;
   TraceOut_MoveRight[132] := BenchUut14.MoveRight;
   TraceOut_ActivateGrip[132] := BenchUut14.ActivateGrip;
   TraceOut_ActivateRelease[132] := BenchUut14.ActivateRelease;
   BenchCalls := BenchCalls + 1;
 133:
   BenchUut14.ManualMode := FALSE;
   BenchUut14.SingleStepMode := TRUE;
   BenchUut14.SingleCycleMode := FALSE;
   BenchUut14.ContinuousMode := FALSE;
   BenchUut14.EmergencyStop := TRUE;
   BenchUut14.Start := FALSE;
   BenchUut14.DownButton := FALSE;
   BenchUut14.UpButton := FALSE;
   BenchUut14.LeftButton := FALSE;
   BenchUut14.RightButton := FALSE;
   BenchUut14.GripButton := FALSE;
   BenchUut14.ReleaseButton := FALSE;
   BenchUut14.DownLimitSwitch := FALSE;
   BenchUut14.UpLimitSwitch := FALSE;
   BenchUut14.LeftLimitSwitch := FALSE;
   BenchUut14.RightLimitSwitch := FALSE;
   BenchUut14.GripLimitSwitch := FALSE;
   BenchUut14.ReleaseLimitSwitch := FALSE;
   TraceIn_ManualMode[133] := BenchUut14.ManualMode;
   TraceIn_SingleStepMode[133] := BenchUut14.SingleStepMode;
   TraceIn_SingleCycleMode[133] := BenchUut14.SingleCycleMode;
   TraceIn_ContinuousMode[133] := BenchUut14.ContinuousMode;
   TraceIn_EmergencyStop[133] := BenchUut14.EmergencyStop;
   TraceIn_Start[133] := BenchUut14.Start;
   TraceIn_DownButton[133] := BenchUut14.DownButton;
   TraceIn_UpButton[133] := BenchUut14.UpButton;
   TraceIn_LeftButton[133] := BenchUut14.LeftButton;
   TraceIn_RightButton[133] := BenchUut14.RightButton;
   TraceIn_GripButton[133] := BenchUut14.GripButton;
   TraceIn_ReleaseButton[133] := BenchUut14.ReleaseButton;
   TraceIn_DownLimitSwitch[133] := BenchUut14.DownLimitSwitch;
   TraceIn_UpLimitSwitch[133] := BenchUut14.UpLimitSwitch;
   TraceIn_LeftLimitSwitch[133] := BenchUut14.LeftLimitSwitch;
   TraceIn_RightLimitSwitch[133] := BenchUut14.RightLimitSwitch;
   TraceIn_GripLimitSwitch[133] := BenchUut14.GripLimitSwitch;
   TraceIn_ReleaseLimitSwitch[133] := BenchUut14.ReleaseLimitSwitch;
   BenchUut14();
   TraceOut_MoveDown[133] := BenchUut14.MoveDown;
   TraceOut_MoveUp[133] := BenchUut14.MoveUp;
   TraceOut_MoveLeft[133] := BenchUut14.MoveLeft;
   TraceOut_MoveRight[133] := BenchUut14.MoveRight;
   TraceOut_ActivateGrip[133] := BenchUut14.ActivateGrip;
   TraceOut_ActivateRelease[133] := BenchUut14.ActivateRelease;
   BenchCalls := BenchCalls + 1;
 134:
   BenchUut14.ManualMode := FALSE;
   BenchUut14.SingleStepMode := TRUE;
   BenchUut14.SingleCycleMode := FALSE;
   BenchUut14.ContinuousMode := FALSE;
   BenchUut14.EmergencyStop := TRUE;
   BenchUut14.Start := FALSE;
   BenchUut14.DownButton := FALSE;
   BenchUut14.UpButton := FALSE;
   BenchUut14.LeftButton := FALSE;
   BenchUut14.RightButton := FALSE;
   BenchUut14.GripButton := FALSE;
   BenchUut14.ReleaseButton := FALSE;
   BenchUut14.DownLimitSwitch := FALSE;
   BenchUut14.UpLimitSwitch := FALSE;
   BenchUut14.LeftLimitSwitch := FALSE;
   BenchUut14.RightLimitSwitch := FALSE;
   BenchUut14.GripLimitSwitch := FALSE;
   BenchUut14.ReleaseLimitSwitch := FALSE;
   TraceIn_ManualMode[134] := BenchUut14.ManualMode;
   TraceIn_SingleStepMode[134] := BenchUut14.SingleStepMode;
   TraceIn_SingleCycleMode[134] := BenchUut14.SingleCycleMode;
   TraceIn_ContinuousMode[134] := BenchUut14.ContinuousMode;
   TraceIn_EmergencyStop[134] := BenchUut14.EmergencyStop;
   TraceIn_Start[134] := BenchUut14.Start;
   TraceIn_DownButton[134] := BenchUut14.DownButton;
   TraceIn_UpButton[134] := BenchUut14.UpButton;
   TraceIn_LeftButton[134] := BenchUut14.LeftButton;
   TraceIn_RightButton[134] := BenchUut14.RightButton;
   TraceIn_GripButton[134] := BenchUut14.GripButton;
   TraceIn_ReleaseButton[134] := BenchUut14.ReleaseButton;
   TraceIn_DownLimitSwitch[134] := BenchUut14.DownLimitSwitch;
   TraceIn_UpLimitSwitch[134] := BenchUut14.UpLimitSwitch;
   TraceIn_LeftLimitSwitch[134] := BenchUut14.LeftLimitSwitch;
   TraceIn_RightLimitSwitch[134] := BenchUut14.RightLimitSwitch;
   TraceIn_GripLimitSwitch[134] := BenchUut14.GripLimitSwitch;
   TraceIn_ReleaseLimitSwitch[134] := BenchUut14.ReleaseLimitSwitch;
   BenchUut14();
   TraceOut_MoveDown[134] := BenchUut14.MoveDown;
   TraceOut_MoveUp[134] := BenchUut14.MoveUp;
   TraceOut_MoveLeft[134] := BenchUut14.MoveLeft;
   TraceOut_MoveRight[134] := BenchUut14.MoveRight;
   TraceOut_ActivateGrip[134] := BenchUut14.ActivateGrip;
   TraceOut_ActivateRelease[134] := BenchUut14.ActivateRelease;
   BenchCalls := BenchCalls + 1;
 135:
   BenchUut14.ManualMode := FALSE;
   BenchUut14.SingleStepMode := TRUE;
   BenchUut14.SingleCycleMode := FALSE;
   BenchUut14.ContinuousMode := FALSE;
   BenchUut14.EmergencyStop := TRUE;
   BenchUut14.Start := FALSE;
   BenchUut14.DownButton := FALSE;
   BenchUut14.UpButton := FALSE;
   BenchUut14.LeftButton := FALSE;
   BenchUut14.RightButton := FALSE;
   BenchUut14.GripButton := FALSE;
   BenchUut14.ReleaseButton := FALSE;
   BenchUut14.DownLimitSwitch := FALSE;
   BenchUut14.UpLimitSwitch := FALSE;
   BenchUut14.LeftLimitSwitch := FALSE;
   BenchUut14.RightLimitSwitch := FALSE;
   BenchUut14.GripLimitSwitch := FALSE;
   BenchUut14.ReleaseLimitSwitch := TRUE;
   TraceIn_ManualMode[135] := BenchUut14.ManualMode;
   TraceIn_SingleStepMode[135] := BenchUut14.SingleStepMode;
   TraceIn_SingleCycleMode[135] := BenchUut14.SingleCycleMode;
   TraceIn_ContinuousMode[135] := BenchUut14.ContinuousMode;
   TraceIn_EmergencyStop[135] := BenchUut14.EmergencyStop;
   TraceIn_Start[135] := BenchUut14.Start;
   TraceIn_DownButton[135] := BenchUut14.DownButton;
   TraceIn_UpButton[135] := BenchUut14.UpButton;
   TraceIn_LeftButton[135] := BenchUut14.LeftButton;
   TraceIn_RightButton[135] := BenchUut14.RightButton;
   TraceIn_GripButton[135] := BenchUut14.GripButton;
   TraceIn_ReleaseButton[135] := BenchUut14.ReleaseButton;
   TraceIn_DownLimitSwitch[135] := BenchUut14.DownLimitSwitch;
   TraceIn_UpLimitSwitch[135] := BenchUut14.UpLimitSwitch;
   TraceIn_LeftLimitSwitch[135] := BenchUut14.LeftLimitSwitch;
   TraceIn_RightLimitSwitch[135] := BenchUut14.RightLimitSwitch;
   TraceIn_GripLimitSwitch[135] := BenchUut14.GripLimitSwitch;
   TraceIn_ReleaseLimitSwitch[135] := BenchUut14.ReleaseLimitSwitch;
   BenchUut14();
   TraceOut_MoveDown[135] := BenchUut14.MoveDown;
   TraceOut_MoveUp[135] := BenchUut14.MoveUp;
   TraceOut_MoveLeft[135] := BenchUut14.MoveLeft;
   TraceOut_MoveRight[135] := BenchUut14.MoveRight;
   TraceOut_ActivateGrip[135] := BenchUut14.ActivateGrip;
   TraceOut_ActivateRelease[135] := BenchUut14.ActivateRelease;
   BenchCalls := BenchCalls + 1;
 136:
   BenchUut14.ManualMode := FALSE;
   BenchUut14.SingleStepMode := TRUE;
   BenchUut14.SingleCycleMode := FALSE;
   BenchUut14.ContinuousMode := FALSE;
   BenchUut14.EmergencyStop := TRUE;
   BenchUut14.Start := TRUE;
   BenchUut14.DownButton := FALSE;
   BenchUut14.UpButton := FALSE;
   BenchUut14.LeftButton := FALSE;
   BenchUut14.RightButton := FALSE;
   BenchUut14.GripButton := FALSE;
   BenchUut14.ReleaseButton := FALSE;
   BenchUut14.DownLimitSwitch := FALSE;
   BenchUut14.UpLimitSwitch := FALSE;
   BenchUut14.LeftLimitSwitch := FALSE;
   BenchUut14.RightLimitSwitch := FALSE;
   BenchUut14.GripLimitSwitch := FALSE;
   BenchUut14.ReleaseLimitSwitch := FALSE;
   TraceIn_ManualMode[136] := BenchUut14.ManualMode;
   TraceIn_SingleStepMode[136] := BenchUut14.SingleStepMode;
   TraceIn_SingleCycleMode[136] := BenchUut14.SingleCycleMode;
   TraceIn_ContinuousMode[136] := BenchUut14.ContinuousMode;
   TraceIn_EmergencyStop[136] := BenchUut14.EmergencyStop;
   TraceIn_Start[136] := BenchUut14.Start;
   TraceIn_DownButton[136] := BenchUut14.DownButton;
   TraceIn_UpButton[136] := BenchUut14.UpButton;
   TraceIn_LeftButton[136] := BenchUut14.LeftButton;
   TraceIn_RightButton[136] := BenchUut14.RightButton;
   TraceIn_GripButton[136] := BenchUut14.GripButton;
   TraceIn_ReleaseButton[136] := BenchUut14.ReleaseButton;
   TraceIn_DownLimitSwitch[136] := BenchUut14.DownLimitSwitch;
   TraceIn_UpLimitSwitch[136] := BenchUut14.UpLimitSwitch;
   TraceIn_LeftLimitSwitch[136] := BenchUut14.LeftLimitSwitch;
   TraceIn_RightLimitSwitch[136] := BenchUut14.RightLimitSwitch;
   TraceIn_GripLimitSwitch[136] := BenchUut14.GripLimitSwitch;
   TraceIn_ReleaseLimitSwitch[136] := BenchUut14.ReleaseLimitSwitch;
   BenchUut14();
   TraceOut_MoveDown[136] := BenchUut14.MoveDown;
   TraceOut_MoveUp[136] := BenchUut14.MoveUp;
   TraceOut_MoveLeft[136] := BenchUut14.MoveLeft;
   TraceOut_MoveRight[136] := BenchUut14.MoveRight;
   TraceOut_ActivateGrip[136] := BenchUut14.ActivateGrip;
   TraceOut_ActivateRelease[136] := BenchUut14.ActivateRelease;
   BenchCalls := BenchCalls + 1;
 137:
   BenchUut14.ManualMode := FALSE;
   BenchUut14.SingleStepMode := TRUE;
   BenchUut14.SingleCycleMode := FALSE;
   BenchUut14.ContinuousMode := FALSE;
   BenchUut14.EmergencyStop := TRUE;
   BenchUut14.Start := FALSE;
   BenchUut14.DownButton := FALSE;
   BenchUut14.UpButton := FALSE;
   BenchUut14.LeftButton := FALSE;
   BenchUut14.RightButton := FALSE;
   BenchUut14.GripButton := FALSE;
   BenchUut14.ReleaseButton := FALSE;
   BenchUut14.DownLimitSwitch := FALSE;
   BenchUut14.UpLimitSwitch := FALSE;
   BenchUut14.LeftLimitSwitch := FALSE;
   BenchUut14.RightLimitSwitch := FALSE;
   BenchUut14.GripLimitSwitch := FALSE;
   BenchUut14.ReleaseLimitSwitch := FALSE;
   TraceIn_ManualMode[137] := BenchUut14.ManualMode;
   TraceIn_SingleStepMode[137] := BenchUut14.SingleStepMode;
   TraceIn_SingleCycleMode[137] := BenchUut14.SingleCycleMode;
   TraceIn_ContinuousMode[137] := BenchUut14.ContinuousMode;
   TraceIn_EmergencyStop[137] := BenchUut14.EmergencyStop;
   TraceIn_Start[137] := BenchUut14.Start;
   TraceIn_DownButton[137] := BenchUut14.DownButton;
   TraceIn_UpButton[137] := BenchUut14.UpButton;
   TraceIn_LeftButton[137] := BenchUut14.LeftButton;
   TraceIn_RightButton[137] := BenchUut14.RightButton;
   TraceIn_GripButton[137] := BenchUut14.GripButton;
   TraceIn_ReleaseButton[137] := BenchUut14.ReleaseButton;
   TraceIn_DownLimitSwitch[137] := BenchUut14.DownLimitSwitch;
   TraceIn_UpLimitSwitch[137] := BenchUut14.UpLimitSwitch;
   TraceIn_LeftLimitSwitch[137] := BenchUut14.LeftLimitSwitch;
   TraceIn_RightLimitSwitch[137] := BenchUut14.RightLimitSwitch;
   TraceIn_GripLimitSwitch[137] := BenchUut14.GripLimitSwitch;
   TraceIn_ReleaseLimitSwitch[137] := BenchUut14.ReleaseLimitSwitch;
   BenchUut14();
   TraceOut_MoveDown[137] := BenchUut14.MoveDown;
   TraceOut_MoveUp[137] := BenchUut14.MoveUp;
   TraceOut_MoveLeft[137] := BenchUut14.MoveLeft;
   TraceOut_MoveRight[137] := BenchUut14.MoveRight;
   TraceOut_ActivateGrip[137] := BenchUut14.ActivateGrip;
   TraceOut_ActivateRelease[137] := BenchUut14.ActivateRelease;
   BenchCalls := BenchCalls + 1;
 138:
   BenchUut14.ManualMode := FALSE;
   BenchUut14.SingleStepMode := TRUE;
   BenchUut14.SingleCycleMode := FALSE;
   BenchUut14.ContinuousMode := FALSE;
   BenchUut14.EmergencyStop := TRUE;
   BenchUut14.Start := FALSE;
   BenchUut14.DownButton := FALSE;
   BenchUut14.UpButton := FALSE;
   BenchUut14.LeftButton := FALSE;
   BenchUut14.RightButton := FALSE;
   BenchUut14.GripButton := FALSE;
   BenchUut14.ReleaseButton := FALSE;
   BenchUut14.DownLimitSwitch := FALSE;
   BenchUut14.UpLimitSwitch := FALSE;
   BenchUut14.LeftLimitSwitch := FALSE;
   BenchUut14.RightLimitSwitch := FALSE;
   BenchUut14.GripLimitSwitch := FALSE;
   BenchUut14.ReleaseLimitSwitch := FALSE;
   TraceIn_ManualMode[138] := BenchUut14.ManualMode;
   TraceIn_SingleStepMode[138] := BenchUut14.SingleStepMode;
   TraceIn_SingleCycleMode[138] := BenchUut14.SingleCycleMode;
   TraceIn_ContinuousMode[138] := BenchUut14.ContinuousMode;
   TraceIn_EmergencyStop[138] := BenchUut14.EmergencyStop;
   TraceIn_Start[138] := BenchUut14.Start;
   TraceIn_DownButton[138] := BenchUut14.DownButton;
   TraceIn_UpButton[138] := BenchUut14.UpButton;
   TraceIn_LeftButton[138] := BenchUut14.LeftButton;
   TraceIn_RightButton[138] := BenchUut14.RightButton;
   TraceIn_GripButton[138] := BenchUut14.GripButton;
   TraceIn_ReleaseButton[138] := BenchUut14.ReleaseButton;
   TraceIn_DownLimitSwitch[138] := BenchUut14.DownLimitSwitch;
   TraceIn_UpLimitSwitch[138] := BenchUut14.UpLimitSwitch;
   TraceIn_LeftLimitSwitch[138] := BenchUut14.LeftLimitSwitch;
   TraceIn_RightLimitSwitch[138] := BenchUut14.RightLimitSwitch;
   TraceIn_GripLimitSwitch[138] := BenchUut14.GripLimitSwitch;
   TraceIn_ReleaseLimitSwitch[138] := BenchUut14.ReleaseLimitSwitch;
   BenchUut14();
   TraceOut_MoveDown[138] := BenchUut14.MoveDown;
   TraceOut_MoveUp[138] := BenchUut14.MoveUp;
   TraceOut_MoveLeft[138] := BenchUut14.MoveLeft;
   TraceOut_MoveRight[138] := BenchUut14.MoveRight;
   TraceOut_ActivateGrip[138] := BenchUut14.ActivateGrip;
   TraceOut_ActivateRelease[138] := BenchUut14.ActivateRelease;
   BenchCalls := BenchCalls + 1;
 139:
   BenchUut14.ManualMode := FALSE;
   BenchUut14.SingleStepMode := TRUE;
   BenchUut14.SingleCycleMode := FALSE;
   BenchUut14.ContinuousMode := FALSE;
   BenchUut14.EmergencyStop := TRUE;
   BenchUut14.Start := FALSE;
   BenchUut14.DownButton := FALSE;
   BenchUut14.UpButton := FALSE;
   BenchUut14.LeftButton := FALSE;
   BenchUut14.RightButton := FALSE;
   BenchUut14.GripButton := FALSE;
   BenchUut14.ReleaseButton := FALSE;
   BenchUut14.DownLimitSwitch := FALSE;
   BenchUut14.UpLimitSwitch := TRUE;
   BenchUut14.LeftLimitSwitch := FALSE;
   BenchUut14.RightLimitSwitch := FALSE;
   BenchUut14.GripLimitSwitch := FALSE;
   BenchUut14.ReleaseLimitSwitch := FALSE;
   TraceIn_ManualMode[139] := BenchUut14.ManualMode;
   TraceIn_SingleStepMode[139] := BenchUut14.SingleStepMode;
   TraceIn_SingleCycleMode[139] := BenchUut14.SingleCycleMode;
   TraceIn_ContinuousMode[139] := BenchUut14.ContinuousMode;
   TraceIn_EmergencyStop[139] := BenchUut14.EmergencyStop;
   TraceIn_Start[139] := BenchUut14.Start;
   TraceIn_DownButton[139] := BenchUut14.DownButton;
   TraceIn_UpButton[139] := BenchUut14.UpButton;
   TraceIn_LeftButton[139] := BenchUut14.LeftButton;
   TraceIn_RightButton[139] := BenchUut14.RightButton;
   TraceIn_GripButton[139] := BenchUut14.GripButton;
   TraceIn_ReleaseButton[139] := BenchUut14.ReleaseButton;
   TraceIn_DownLimitSwitch[139] := BenchUut14.DownLimitSwitch;
   TraceIn_UpLimitSwitch[139] := BenchUut14.UpLimitSwitch;
   TraceIn_LeftLimitSwitch[139] := BenchUut14.LeftLimitSwitch;
   TraceIn_RightLimitSwitch[139] := BenchUut14.RightLimitSwitch;
   TraceIn_GripLimitSwitch[139] := BenchUut14.GripLimitSwitch;
   TraceIn_ReleaseLimitSwitch[139] := BenchUut14.ReleaseLimitSwitch;
   BenchUut14();
   TraceOut_MoveDown[139] := BenchUut14.MoveDown;
   TraceOut_MoveUp[139] := BenchUut14.MoveUp;
   TraceOut_MoveLeft[139] := BenchUut14.MoveLeft;
   TraceOut_MoveRight[139] := BenchUut14.MoveRight;
   TraceOut_ActivateGrip[139] := BenchUut14.ActivateGrip;
   TraceOut_ActivateRelease[139] := BenchUut14.ActivateRelease;
   BenchCalls := BenchCalls + 1;
 140:
   BenchUut14.ManualMode := FALSE;
   BenchUut14.SingleStepMode := TRUE;
   BenchUut14.SingleCycleMode := FALSE;
   BenchUut14.ContinuousMode := FALSE;
   BenchUut14.EmergencyStop := TRUE;
   BenchUut14.Start := TRUE;
   BenchUut14.DownButton := FALSE;
   BenchUut14.UpButton := FALSE;
   BenchUut14.LeftButton := FALSE;
   BenchUut14.RightButton := FALSE;
   BenchUut14.GripButton := FALSE;
   BenchUut14.ReleaseButton := FALSE;
   BenchUut14.DownLimitSwitch := FALSE;
   BenchUut14.UpLimitSwitch := FALSE;
   BenchUut14.LeftLimitSwitch := FALSE;
   BenchUut14.RightLimitSwitch := FALSE;
   BenchUut14.GripLimitSwitch := FALSE;
   BenchUut14.ReleaseLimitSwitch := FALSE;
   TraceIn_ManualMode[140] := BenchUut14.ManualMode;
   TraceIn_SingleStepMode[140] := BenchUut14.SingleStepMode;
   TraceIn_SingleCycleMode[140] := BenchUut14.SingleCycleMode;
   TraceIn_ContinuousMode[140] := BenchUut14.ContinuousMode;
   TraceIn_EmergencyStop[140] := BenchUut14.EmergencyStop;
   TraceIn_Start[140] := BenchUut14.Start;
   TraceIn_DownButton[140] := BenchUut14.DownButton;
   TraceIn_UpButton[140] := BenchUut14.UpButton;
   TraceIn_LeftButton[140] := BenchUut14.LeftButton;
   TraceIn_RightButton[140] := BenchUut14.RightButton;
   TraceIn_GripButton[140] := BenchUut14.GripButton;
   TraceIn_ReleaseButton[140] := BenchUut14.ReleaseButton;
   TraceIn_DownLimitSwitch[140] := BenchUut14.DownLimitSwitch;
   TraceIn_UpLimitSwitch[140] := BenchUut14.UpLimitSwitch;
   TraceIn_LeftLimitSwitch[140] := BenchUut14.LeftLimitSwitch;
   TraceIn_RightLimitSwitch[140] := BenchUut14.RightLimitSwitch;
   TraceIn_GripLimitSwitch[140] := BenchUut14.GripLimitSwitch;
   TraceIn_ReleaseLimitSwitch[140] := BenchUut14.ReleaseLimitSwitch;
   BenchUut14();
   TraceOut_MoveDown[140] := BenchUut14.MoveDown;
   TraceOut_MoveUp[140] := BenchUut14.MoveUp;
   TraceOut_MoveLeft[140] := BenchUut14.MoveLeft;
   TraceOut_MoveRight[140] := BenchUut14.MoveRight;
   TraceOut_ActivateGrip[140] := BenchUut14.ActivateGrip;
   TraceOut_ActivateRelease[140] := BenchUut14.ActivateRelease;
   BenchCalls := BenchCalls + 1;
 141:
   BenchUut14.ManualMode := FALSE;
   BenchUut14.SingleStepMode := TRUE;
   BenchUut14.SingleCycleMode := FALSE;
   BenchUut14.ContinuousMode := FALSE;
   BenchUut14.EmergencyStop := TRUE;
   BenchUut14.Start := FALSE;
   BenchUut14.DownButton := FALSE;
   BenchUut14.UpButton := FALSE;
   BenchUut14.LeftButton := FALSE;
   BenchUut14.RightButton := FALSE;
   BenchUut14.GripButton := FALSE;
   BenchUut14.ReleaseButton := FALSE;
   BenchUut14.DownLimitSwitch := FALSE;
   BenchUut14.UpLimitSwitch := FALSE;
   BenchUut14.LeftLimitSwitch := FALSE;
   BenchUut14.RightLimitSwitch := FALSE;
   BenchUut14.GripLimitSwitch := FALSE;
   BenchUut14.ReleaseLimitSwitch := FALSE;
   TraceIn_ManualMode[141] := BenchUut14.ManualMode;
   TraceIn_SingleStepMode[141] := BenchUut14.SingleStepMode;
   TraceIn_SingleCycleMode[141] := BenchUut14.SingleCycleMode;
   TraceIn_ContinuousMode[141] := BenchUut14.ContinuousMode;
   TraceIn_EmergencyStop[141] := BenchUut14.EmergencyStop;
   TraceIn_Start[141] := BenchUut14.Start;
   TraceIn_DownButton[141] := BenchUut14.DownButton;
   TraceIn_UpButton[141] := BenchUut14.UpButton;
   TraceIn_LeftButton[141] := BenchUut14.LeftButton;
   TraceIn_RightButton[141] := BenchUut14.RightButton;
   TraceIn_GripButton[141] := BenchUut14.GripButton;
   TraceIn_ReleaseButton[141] := BenchUut14.ReleaseButton;
   TraceIn_DownLimitSwitch[141] := BenchUut14.DownLimitSwitch;
   TraceIn_UpLimitSwitch[141] := BenchUut14.UpLimitSwitch;
   TraceIn_LeftLimitSwitch[141] := BenchUut14.LeftLimitSwitch;
   TraceIn_RightLimitSwitch[141] := BenchUut14.RightLimitSwitch;
   TraceIn_GripLimitSwitch[141] := BenchUut14.GripLimitSwitch;
   TraceIn_ReleaseLimitSwitch[141] := BenchUut14.ReleaseLimitSwitch;
   BenchUut14();
   TraceOut_MoveDown[141] := BenchUut14.MoveDown;
   TraceOut_MoveUp[141] := BenchUut14.MoveUp;
   TraceOut_MoveLeft[141] := BenchUut14.MoveLeft;
   TraceOut_MoveRight[141] := BenchUut14.MoveRight;
   TraceOut_ActivateGrip[141] := BenchUut14.ActivateGrip;
   TraceOut_ActivateRelease[141] := BenchUut14.ActivateRelease;
   BenchCalls := BenchCalls + 1;
 142:
   BenchUut14.ManualMode := FALSE;
   BenchUut14.SingleStepMode := TRUE;
   BenchUut14.SingleCycleMode := FALSE;
   BenchUut14.ContinuousMode := FALSE;
   BenchUut14.EmergencyStop := TRUE;
   BenchUut14.Start := FALSE;
   BenchUut14.DownButton := FALSE;
   BenchUut14.UpButton := FALSE;
   BenchUut14.LeftButton := FALSE;
   BenchUut14.RightButton := FALSE;
   BenchUut14.GripButton := FALSE;
   BenchUut14.ReleaseButton := FALSE;
   BenchUut14.DownLimitSwitch := FALSE;
   BenchUut14.UpLimitSwitch := FALSE;
   BenchUut14.LeftLimitSwitch := FALSE;
   BenchUut14.RightLimitSwitch := FALSE;
   BenchUut14.GripLimitSwitch := FALSE;
   BenchUut14.ReleaseLimitSwitch := FALSE;
   TraceIn_ManualMode[142] := BenchUut14.ManualMode;
   TraceIn_SingleStepMode[142] := BenchUut14.SingleStepMode;
   TraceIn_SingleCycleMode[142] := BenchUut14.SingleCycleMode;
   TraceIn_ContinuousMode[142] := BenchUut14.ContinuousMode;
   TraceIn_EmergencyStop[142] := BenchUut14.EmergencyStop;
   TraceIn_Start[142] := BenchUut14.Start;
   TraceIn_DownButton[142] := BenchUut14.DownButton;
   TraceIn_UpButton[142] := BenchUut14.UpButton;
   TraceIn_LeftButton[142] := BenchUut14.LeftButton;
   TraceIn_RightButton[142] := BenchUut14.RightButton;
   TraceIn_GripButton[142] := BenchUut14.GripButton;
   TraceIn_ReleaseButton[142] := BenchUut14.ReleaseButton;
   TraceIn_DownLimitSwitch[142] := BenchUut14.DownLimitSwitch;
   TraceIn_UpLimitSwitch[142] := BenchUut14.UpLimitSwitch;
   TraceIn_LeftLimitSwitch[142] := BenchUut14.LeftLimitSwitch;
   TraceIn_RightLimitSwitch[142] := BenchUut14.RightLimitSwitch;
   TraceIn_GripLimitSwitch[142] := BenchUut14.GripLimitSwitch;
   TraceIn_ReleaseLimitSwitch[142] := BenchUut14.ReleaseLimitSwitch;
   BenchUut14();
   TraceOut_MoveDown[142] := BenchUut14.MoveDown;
   TraceOut_MoveUp[142] := BenchUut14.MoveUp;
   TraceOut_MoveLeft[142] := BenchUut14.MoveLeft;
   TraceOut_MoveRight[142] := BenchUut14.MoveRight;
   TraceOut_ActivateGrip[142] := BenchUut14.ActivateGrip;
   TraceOut_ActivateRelease[142] := BenchUut14.ActivateRelease;
   BenchCalls := BenchCalls + 1;
 143:
   BenchUut14.ManualMode := FALSE;
   BenchUut14.SingleStepMode := TRUE;
   BenchUut14.SingleCycleMode := FALSE;
   BenchUut14.ContinuousMode := FALSE;
   BenchUut14.EmergencyStop := TRUE;
   BenchUut14.Start := FALSE;
   BenchUut14.DownButton := FALSE;
   BenchUut14.UpButton := FALSE;
   BenchUut14.LeftButton := FALSE;
   BenchUut14.RightButton := FALSE;
   BenchUut14.GripButton := FALSE;
   BenchUut14.ReleaseButton := FALSE;
   BenchUut14.DownLimitSwitch := FALSE;
   BenchUut14.UpLimitSwitch := FALSE;
   BenchUut14.LeftLimitSwitch := TRUE;
   BenchUut14.RightLimitSwitch := FALSE;
   BenchUut14.GripLimitSwitch := FALSE;
   BenchUut14.ReleaseLimitSwitch := FALSE;
   TraceIn_ManualMode[143] := BenchUut14.ManualMode;
   TraceIn_SingleStepMode[143] := BenchUut14.SingleStepMode;
   TraceIn_SingleCycleMode[143] := BenchUut14.SingleCycleMode;
   TraceIn_ContinuousMode[143] := BenchUut14.ContinuousMode;
   TraceIn_EmergencyStop[143] := BenchUut14.EmergencyStop;
   TraceIn_Start[143] := BenchUut14.Start;
   TraceIn_DownButton[143] := BenchUut14.DownButton;
   TraceIn_UpButton[143] := BenchUut14.UpButton;
   TraceIn_LeftButton[143] := BenchUut14.LeftButton;
   TraceIn_RightButton[143] := BenchUut14.RightButton;
   TraceIn_GripButton[143] := BenchUut14.GripButton;
   TraceIn_ReleaseButton[143] := BenchUut14.ReleaseButton;
   TraceIn_DownLimitSwitch[143] := BenchUut14.DownLimitSwitch;
   TraceIn_UpLimitSwitch[143] := BenchUut14.UpLimitSwitch;
   TraceIn_LeftLimitSwitch[143] := BenchUut14.LeftLimitSwitch;
   TraceIn_RightLimitSwitch[143] := BenchUut14.RightLimitSwitch;
   TraceIn_GripLimitSwitch[143] := BenchUut14.GripLimitSwitch;
   TraceIn_ReleaseLimitSwitch[143] := BenchUut14.ReleaseLimitSwitch;
   BenchUut14();
   TraceOut_MoveDown[143] := BenchUut14.MoveDown;
   TraceOut_MoveUp[143] := BenchUut14.MoveUp;
   TraceOut_MoveLeft[143] := BenchUut14.MoveLeft;
   TraceOut_MoveRight[143] := BenchUut14.MoveRight;
   TraceOut_ActivateGrip[143] := BenchUut14.ActivateGrip;
   TraceOut_ActivateRelease[143] := BenchUut14.ActivateRelease;
   BenchCalls := BenchCalls + 1;
 144:
   BenchUut14.ManualMode := FALSE;
   BenchUut14.SingleStepMode := TRUE;
   BenchUut14.SingleCycleMode := FALSE;
   BenchUut14.ContinuousMode := FALSE;
   BenchUut14.EmergencyStop := TRUE;
   BenchUut14.Start := TRUE;
   BenchUut14.DownButton := FALSE;
   BenchUut14.UpButton := FALSE;
   BenchUut14.LeftButton := FALSE;
   BenchUut14.RightButton := FALSE;
   BenchUut14.GripButton := FALSE;
   BenchUut14.ReleaseButton := FALSE;
   BenchUut14.DownLimitSwitch := FALSE;
   BenchUut14.UpLimitSwitch := TRUE;
   BenchUut14.LeftLimitSwitch := TRUE;
   BenchUut14.RightLimitSwitch := FALSE;
   BenchUut14.GripLimitSwitch := FALSE;
   BenchUut14.ReleaseLimitSwitch := FALSE;
   TraceIn_ManualMode[144] := BenchUut14.ManualMode;
   TraceIn_SingleStepMode[144] := BenchUut14.SingleStepMode;
   TraceIn_SingleCycleMode[144] := BenchUut14.SingleCycleMode;
   TraceIn_ContinuousMode[144] := BenchUut14.ContinuousMode;
   TraceIn_EmergencyStop[144] := BenchUut14.EmergencyStop;
   TraceIn_Start[144] := BenchUut14.Start;
   TraceIn_DownButton[144] := BenchUut14.DownButton;
   TraceIn_UpButton[144] := BenchUut14.UpButton;
   TraceIn_LeftButton[144] := BenchUut14.LeftButton;
   TraceIn_RightButton[144] := BenchUut14.RightButton;
   TraceIn_GripButton[144] := BenchUut14.GripButton;
   TraceIn_ReleaseButton[144] := BenchUut14.ReleaseButton;
   TraceIn_DownLimitSwitch[144] := BenchUut14.DownLimitSwitch;
   TraceIn_UpLimitSwitch[144] := BenchUut14.UpLimitSwitch;
   TraceIn_LeftLimitSwitch[144] := BenchUut14.LeftLimitSwitch;
   TraceIn_RightLimitSwitch[144] := BenchUut14.RightLimitSwitch;
   TraceIn_GripLimitSwitch[144] := BenchUut14.GripLimitSwitch;
   TraceIn_ReleaseLimitSwitch[144] := BenchUut14.ReleaseLimitSwitch;
   BenchUut14();
   TraceOut_MoveDown[144] := BenchUut14.MoveDown;
   TraceOut_MoveUp[144] := BenchUut14.MoveUp;
   TraceOut_MoveLeft[144] := BenchUut14.MoveLeft;
   TraceOut_MoveRight[144] := BenchUut14.MoveRight;
   TraceOut_ActivateGrip[144] := BenchUut14.ActivateGrip;
   TraceOut_ActivateRelease[144] := BenchUut14.ActivateRelease;
   BenchCalls := BenchCalls + 1;
 145:
   BenchUut14.ManualMode := FALSE;
   BenchUut14.SingleStepMode := TRUE;
   BenchUut14.SingleCycleMode := FALSE;
   BenchUut14.ContinuousMode := FALSE;
   BenchUut14.EmergencyStop := TRUE;
   BenchUut14.Start := FALSE;
   BenchUut14.DownButton := FALSE;
   BenchUut14.UpButton := FALSE;
   BenchUut14.LeftButton := FALSE;
   BenchUut14.RightButton := FALSE;
   BenchUut14.GripButton := FALSE;
   BenchUut14.ReleaseButton := FALSE;
   BenchUut14.DownLimitSwitch := FALSE;
   BenchUut14.UpLimitSwitch := TRUE;
   BenchUut14.LeftLimitSwitch := TRUE;
   BenchUut14.RightLimitSwitch := FALSE;
   BenchUut14.GripLimitSwitch := FALSE;
   BenchUut14.ReleaseLimitSwitch := FALSE;
   TraceIn_ManualMode[145] := BenchUut14.ManualMode;
   TraceIn_SingleStepMode[145] := BenchUut14.SingleStepMode;
   TraceIn_SingleCycleMode[145] := BenchUut14.SingleCycleMode;
   TraceIn_ContinuousMode[145] := BenchUut14.ContinuousMode;
   TraceIn_EmergencyStop[145] := BenchUut14.EmergencyStop;
   TraceIn_Start[145] := BenchUut14.Start;
   TraceIn_DownButton[145] := BenchUut14.DownButton;
   TraceIn_UpButton[145] := BenchUut14.UpButton;
   TraceIn_LeftButton[145] := BenchUut14.LeftButton;
   TraceIn_RightButton[145] := BenchUut14.RightButton;
   TraceIn_GripButton[145] := BenchUut14.GripButton;
   TraceIn_ReleaseButton[145] := BenchUut14.ReleaseButton;
   TraceIn_DownLimitSwitch[145] := BenchUut14.DownLimitSwitch;
   TraceIn_UpLimitSwitch[145] := BenchUut14.UpLimitSwitch;
   TraceIn_LeftLimitSwitch[145] := BenchUut14.LeftLimitSwitch;
   TraceIn_RightLimitSwitch[145] := BenchUut14.RightLimitSwitch;
   TraceIn_GripLimitSwitch[145] := BenchUut14.GripLimitSwitch;
   TraceIn_ReleaseLimitSwitch[145] := BenchUut14.ReleaseLimitSwitch;
   BenchUut14();
   TraceOut_MoveDown[145] := BenchUut14.MoveDown;
   TraceOut_MoveUp[145] := BenchUut14.MoveUp;
   TraceOut_MoveLeft[145] := BenchUut14.MoveLeft;
   TraceOut_MoveRight[145] := BenchUut14.MoveRight;
   TraceOut_ActivateGrip[145] := BenchUut14.ActivateGrip;
   TraceOut_ActivateRelease[145] := BenchUut14.ActivateRelease;
   BenchCalls := BenchCalls + 1;
 146:
   BenchUut14.ManualMode := FALSE;
   BenchUut14.SingleStepMode := TRUE;
   BenchUut14.SingleCycleMode := FALSE;
   BenchUut14.ContinuousMode := FALSE;
   BenchUut14.EmergencyStop := TRUE;
   BenchUut14.Start := FALSE;
   BenchUut14.DownButton := FALSE;
   BenchUut14.UpButton := FALSE;
   BenchUut14.LeftButton := FALSE;
   BenchUut14.RightButton := FALSE;
   BenchUut14.GripButton := FALSE;
   BenchUut14.ReleaseButton := FALSE;
   BenchUut14.DownLimitSwitch := FALSE;
   BenchUut14.UpLimitSwitch := TRUE;
   BenchUut14.LeftLimitSwitch := TRUE;
   BenchUut14.RightLimitSwitch := FALSE;
   BenchUut14.GripLimitSwitch := FALSE;
   BenchUut14.ReleaseLimitSwitch := FALSE;
   TraceIn_ManualMode[146] := BenchUut14.ManualMode;
   TraceIn_SingleStepMode[146] := BenchUut14.SingleStepMode;
   TraceIn_SingleCycleMode[146] := BenchUut14.SingleCycleMode;
   TraceIn_ContinuousMode[146] := BenchUut14.ContinuousMode;
   TraceIn_EmergencyStop[146] := BenchUut14.EmergencyStop;
   TraceIn_Start[146] := BenchUut14.Start;
   TraceIn_DownButton[146] := BenchUut14.DownButton;
   TraceIn_UpButton[146] := BenchUut14.UpButton;
   TraceIn_LeftButton[146] := BenchUut14.LeftButton;
   TraceIn_RightButton[146] := BenchUut14.RightButton;
   TraceIn_GripButton[146] := BenchUut14.GripButton;
   TraceIn_ReleaseButton[146] := BenchUut14.ReleaseButton;
   TraceIn_DownLimitSwitch[146] := BenchUut14.DownLimitSwitch;
   TraceIn_UpLimitSwitch[146] := BenchUut14.UpLimitSwitch;
   TraceIn_LeftLimitSwitch[146] := BenchUut14.LeftLimitSwitch;
   TraceIn_RightLimitSwitch[146] := BenchUut14.RightLimitSwitch;
   TraceIn_GripLimitSwitch[146] := BenchUut14.GripLimitSwitch;
   TraceIn_ReleaseLimitSwitch[146] := BenchUut14.ReleaseLimitSwitch;
   BenchUut14();
   TraceOut_MoveDown[146] := BenchUut14.MoveDown;
   TraceOut_MoveUp[146] := BenchUut14.MoveUp;
   TraceOut_MoveLeft[146] := BenchUut14.MoveLeft;
   TraceOut_MoveRight[146] := BenchUut14.MoveRight;
   TraceOut_ActivateGrip[146] := BenchUut14.ActivateGrip;
   TraceOut_ActivateRelease[146] := BenchUut14.ActivateRelease;
   BenchCalls := BenchCalls + 1;
 147:
   BenchUut14.ManualMode := FALSE;
   BenchUut14.SingleStepMode := TRUE;
   BenchUut14.SingleCycleMode := FALSE;
   BenchUut14.ContinuousMode := FALSE;
   BenchUut14.EmergencyStop := TRUE;
   BenchUut14.Start := FALSE;
   BenchUut14.DownButton := FALSE;
   BenchUut14.UpButton := FALSE;
   BenchUut14.LeftButton := FALSE;
   BenchUut14.RightButton := FALSE;
   BenchUut14.GripButton := FALSE;
   BenchUut14.ReleaseButton := FALSE;
   BenchUut14.DownLimitSwitch := TRUE;
   BenchUut14.UpLimitSwitch := FALSE;
   BenchUut14.LeftLimitSwitch := FALSE;
   BenchUut14.RightLimitSwitch := FALSE;
   BenchUut14.GripLimitSwitch := FALSE;
   BenchUut14.ReleaseLimitSwitch := FALSE;
   TraceIn_ManualMode[147] := BenchUut14.ManualMode;
   TraceIn_SingleStepMode[147] := BenchUut14.SingleStepMode;
   TraceIn_SingleCycleMode[147] := BenchUut14.SingleCycleMode;
   TraceIn_ContinuousMode[147] := BenchUut14.ContinuousMode;
   TraceIn_EmergencyStop[147] := BenchUut14.EmergencyStop;
   TraceIn_Start[147] := BenchUut14.Start;
   TraceIn_DownButton[147] := BenchUut14.DownButton;
   TraceIn_UpButton[147] := BenchUut14.UpButton;
   TraceIn_LeftButton[147] := BenchUut14.LeftButton;
   TraceIn_RightButton[147] := BenchUut14.RightButton;
   TraceIn_GripButton[147] := BenchUut14.GripButton;
   TraceIn_ReleaseButton[147] := BenchUut14.ReleaseButton;
   TraceIn_DownLimitSwitch[147] := BenchUut14.DownLimitSwitch;
   TraceIn_UpLimitSwitch[147] := BenchUut14.UpLimitSwitch;
   TraceIn_LeftLimitSwitch[147] := BenchUut14.LeftLimitSwitch;
   TraceIn_RightLimitSwitch[147] := BenchUut14.RightLimitSwitch;
   TraceIn_GripLimitSwitch[147] := BenchUut14.GripLimitSwitch;
   TraceIn_ReleaseLimitSwitch[147] := BenchUut14.ReleaseLimitSwitch;
   BenchUut14();
   TraceOut_MoveDown[147] := BenchUut14.MoveDown;
   TraceOut_MoveUp[147] := BenchUut14.MoveUp;
   TraceOut_MoveLeft[147] := BenchUut14.MoveLeft;
   TraceOut_MoveRight[147] := BenchUut14.MoveRight;
   TraceOut_ActivateGrip[147] := BenchUut14.ActivateGrip;
   TraceOut_ActivateRelease[147] := BenchUut14.ActivateRelease;
   BenchCalls := BenchCalls + 1;
 148:
   BenchUut14.ManualMode := FALSE;
   BenchUut14.SingleStepMode := TRUE;
   BenchUut14.SingleCycleMode := FALSE;
   BenchUut14.ContinuousMode := FALSE;
   BenchUut14.EmergencyStop := TRUE;
   BenchUut14.Start := TRUE;
   BenchUut14.DownButton := FALSE;
   BenchUut14.UpButton := FALSE;
   BenchUut14.LeftButton := FALSE;
   BenchUut14.RightButton := FALSE;
   BenchUut14.GripButton := FALSE;
   BenchUut14.ReleaseButton := FALSE;
   BenchUut14.DownLimitSwitch := FALSE;
   BenchUut14.UpLimitSwitch := FALSE;
   BenchUut14.LeftLimitSwitch := FALSE;
   BenchUut14.RightLimitSwitch := FALSE;
   BenchUut14.GripLimitSwitch := FALSE;
   BenchUut14.ReleaseLimitSwitch := FALSE;
   TraceIn_ManualMode[148] := BenchUut14.ManualMode;
   TraceIn_SingleStepMode[148] := BenchUut14.SingleStepMode;
   TraceIn_SingleCycleMode[148] := BenchUut14.SingleCycleMode;
   TraceIn_ContinuousMode[148] := BenchUut14.ContinuousMode;
   TraceIn_EmergencyStop[148] := BenchUut14.EmergencyStop;
   TraceIn_Start[148] := BenchUut14.Start;
   TraceIn_DownButton[148] := BenchUut14.DownButton;
   TraceIn_UpButton[148] := BenchUut14.UpButton;
   TraceIn_LeftButton[148] := BenchUut14.LeftButton;
   TraceIn_RightButton[148] := BenchUut14.RightButton;
   TraceIn_GripButton[148] := BenchUut14.GripButton;
   TraceIn_ReleaseButton[148] := BenchUut14.ReleaseButton;
   TraceIn_DownLimitSwitch[148] := BenchUut14.DownLimitSwitch;
   TraceIn_UpLimitSwitch[148] := BenchUut14.UpLimitSwitch;
   TraceIn_LeftLimitSwitch[148] := BenchUut14.LeftLimitSwitch;
   TraceIn_RightLimitSwitch[148] := BenchUut14.RightLimitSwitch;
   TraceIn_GripLimitSwitch[148] := BenchUut14.GripLimitSwitch;
   TraceIn_ReleaseLimitSwitch[148] := BenchUut14.ReleaseLimitSwitch;
   BenchUut14();
   TraceOut_MoveDown[148] := BenchUut14.MoveDown;
   TraceOut_MoveUp[148] := BenchUut14.MoveUp;
   TraceOut_MoveLeft[148] := BenchUut14.MoveLeft;
   TraceOut_MoveRight[148] := BenchUut14.MoveRight;
   TraceOut_ActivateGrip[148] := BenchUut14.ActivateGrip;
   TraceOut_ActivateRelease[148] := BenchUut14.ActivateRelease;
   BenchCalls := BenchCalls + 1;
 149:
   BenchUut14.ManualMode := FALSE;
   BenchUut14.SingleStepMode := TRUE;
   BenchUut14.SingleCycleMode := FALSE;
   BenchUut14.ContinuousMode := FALSE;
   BenchUut14.EmergencyStop := TRUE;
   BenchUut14.Start := FALSE;
   BenchUut14.DownButton := FALSE;
   BenchUut14.UpButton := FALSE;
   BenchUut14.LeftButton := FALSE;
   BenchUut14.RightButton := FALSE;
   BenchUut14.GripButton := FALSE;
   BenchUut14.ReleaseButton := FALSE;
   BenchUut14.DownLimitSwitch := FALSE;
   BenchUut14.UpLimitSwitch := FALSE;
   BenchUut14.LeftLimitSwitch := FALSE;
   BenchUut14.RightLimitSwitch := FALSE;
   BenchUut14.GripLimitSwitch := FALSE;
   BenchUut14.ReleaseLimitSwitch := FALSE;
   TraceIn_ManualMode[149] := BenchUut14.ManualMode;
   TraceIn_SingleStepMode[149] := BenchUut14.SingleStepMode;
   TraceIn_SingleCycleMode[149] := BenchUut14.SingleCycleMode;
   TraceIn_ContinuousMode[149] := BenchUut14.ContinuousMode;
   TraceIn_EmergencyStop[149] := BenchUut14.EmergencyStop;
   TraceIn_Start[149] := BenchUut14.Start;
   TraceIn_DownButton[149] := BenchUut14.DownButton;
   TraceIn_UpButton[149] := BenchUut14.UpButton;
   TraceIn_LeftButton[149] := BenchUut14.LeftButton;
   TraceIn_RightButton[149] := BenchUut14.RightButton;
   TraceIn_GripButton[149] := BenchUut14.GripButton;
   TraceIn_ReleaseButton[149] := BenchUut14.ReleaseButton;
   TraceIn_DownLimitSwitch[149] := BenchUut14.DownLimitSwitch;
   TraceIn_UpLimitSwitch[149] := BenchUut14.UpLimitSwitch;
   TraceIn_LeftLimitSwitch[149] := BenchUut14.LeftLimitSwitch;
   TraceIn_RightLimitSwitch[149] := BenchUut14.RightLimitSwitch;
   TraceIn_GripLimitSwitch[149] := BenchUut14.GripLimitSwitch;
   TraceIn_ReleaseLimitSwitch[149] := BenchUut14.ReleaseLimitSwitch;
   BenchUut14();
   TraceOut_MoveDown[149] := BenchUut14.MoveDown;
   TraceOut_MoveUp[149] := BenchUut14.MoveUp;
   TraceOut_MoveLeft[149] := BenchUut14.MoveLeft;
   TraceOut_MoveRight[149] := BenchUut14.MoveRight;
   TraceOut_ActivateGrip[149] := BenchUut14.ActivateGrip;
   TraceOut_ActivateRelease[149] := BenchUut14.ActivateRelease;
   BenchCalls := BenchCalls + 1;
 150:
   BenchUut14.ManualMode := FALSE;
   BenchUut14.SingleStepMode := TRUE;
   BenchUut14.SingleCycleMode := FALSE;
   BenchUut14.ContinuousMode := FALSE;
   BenchUut14.EmergencyStop := TRUE;
   BenchUut14.Start := FALSE;
   BenchUut14.DownButton := FALSE;
   BenchUut14.UpButton := FALSE;
   BenchUut14.LeftButton := FALSE;
   BenchUut14.RightButton := FALSE;
   BenchUut14.GripButton := FALSE;
   BenchUut14.ReleaseButton := FALSE;
   BenchUut14.DownLimitSwitch := FALSE;
   BenchUut14.UpLimitSwitch := FALSE;
   BenchUut14.LeftLimitSwitch := FALSE;
   BenchUut14.RightLimitSwitch := FALSE;
   BenchUut14.GripLimitSwitch := FALSE;
   BenchUut14.ReleaseLimitSwitch := FALSE;
   TraceIn_ManualMode[150] := BenchUut14.ManualMode;
   TraceIn_SingleStepMode[150] := BenchUut14.SingleStepMode;
   TraceIn_SingleCycleMode[150] := BenchUut14.SingleCycleMode;
   TraceIn_ContinuousMode[150] := BenchUut14.ContinuousMode;
   TraceIn_EmergencyStop[150] := BenchUut14.EmergencyStop;
   TraceIn_Start[150] := BenchUut14.Start;
   TraceIn_DownButton[150] := BenchUut14.DownButton;
   TraceIn_UpButton[150] := BenchUut14.UpButton;
   TraceIn_LeftButton[150] := BenchUut14.LeftButton;
   TraceIn_RightButton[150] := BenchUut14.RightButton;
   TraceIn_GripButton[150] := BenchUut14.GripButton;
   TraceIn_ReleaseButton[150] := BenchUut14.ReleaseButton;
   TraceIn_DownLimitSwitch[150] := BenchUut14.DownLimitSwitch;
   TraceIn_UpLimitSwitch[150] := BenchUut14.UpLimitSwitch;
   TraceIn_LeftLimitSwitch[150] := BenchUut14.LeftLimitSwitch;
   TraceIn_RightLimitSwitch[150] := BenchUut14.RightLimitSwitch;
   TraceIn_GripLimitSwitch[150] := BenchUut14.GripLimitSwitch;
   TraceIn_ReleaseLimitSwitch[150] := BenchUut14.ReleaseLimitSwitch;
   BenchUut14();
   TraceOut_MoveDown[150] := BenchUut14.MoveDown;
   TraceOut_MoveUp[150] := BenchUut14.MoveUp;
   TraceOut_MoveLeft[150] := BenchUut14.MoveLeft;
   TraceOut_MoveRight[150] := BenchUut14.MoveRight;
   TraceOut_ActivateGrip[150] := BenchUut14.ActivateGrip;
   TraceOut_ActivateRelease[150] := BenchUut14.ActivateRelease;
   BenchCalls := BenchCalls + 1;
 151:
   BenchUut14.ManualMode := FALSE;
   BenchUut14.SingleStepMode := TRUE;
   BenchUut14.SingleCycleMode := FALSE;
   BenchUut14.ContinuousMode := FALSE;
   BenchUut14.EmergencyStop := TRUE;
   BenchUut14.Start := FALSE;
   BenchUut14.DownButton := FALSE;
   BenchUut14.UpButton := FALSE;
   BenchUut14.LeftButton := FALSE;
   BenchUut14.RightButton := FALSE;
   BenchUut14.GripButton := FALSE;
   BenchUut14.ReleaseButton := FALSE;
   BenchUut14.DownLimitSwitch := FALSE;
   BenchUut14.UpLimitSwitch := FALSE;
   BenchUut14.LeftLimitSwitch := FALSE;
   BenchUut14.RightLimitSwitch := FALSE;
   BenchUut14.GripLimitSwitch := TRUE;
   BenchUut14.ReleaseLimitSwitch := FALSE;
   TraceIn_ManualMode[151] := BenchUut14.ManualMode;
   TraceIn_SingleStepMode[151] := BenchUut14.SingleStepMode;
   TraceIn_SingleCycleMode[151] := BenchUut14.SingleCycleMode;
   TraceIn_ContinuousMode[151] := BenchUut14.ContinuousMode;
   TraceIn_EmergencyStop[151] := BenchUut14.EmergencyStop;
   TraceIn_Start[151] := BenchUut14.Start;
   TraceIn_DownButton[151] := BenchUut14.DownButton;
   TraceIn_UpButton[151] := BenchUut14.UpButton;
   TraceIn_LeftButton[151] := BenchUut14.LeftButton;
   TraceIn_RightButton[151] := BenchUut14.RightButton;
   TraceIn_GripButton[151] := BenchUut14.GripButton;
   TraceIn_ReleaseButton[151] := BenchUut14.ReleaseButton;
   TraceIn_DownLimitSwitch[151] := BenchUut14.DownLimitSwitch;
   TraceIn_UpLimitSwitch[151] := BenchUut14.UpLimitSwitch;
   TraceIn_LeftLimitSwitch[151] := BenchUut14.LeftLimitSwitch;
   TraceIn_RightLimitSwitch[151] := BenchUut14.RightLimitSwitch;
   TraceIn_GripLimitSwitch[151] := BenchUut14.GripLimitSwitch;
   TraceIn_ReleaseLimitSwitch[151] := BenchUut14.ReleaseLimitSwitch;
   BenchUut14();
   TraceOut_MoveDown[151] := BenchUut14.MoveDown;
   TraceOut_MoveUp[151] := BenchUut14.MoveUp;
   TraceOut_MoveLeft[151] := BenchUut14.MoveLeft;
   TraceOut_MoveRight[151] := BenchUut14.MoveRight;
   TraceOut_ActivateGrip[151] := BenchUut14.ActivateGrip;
   TraceOut_ActivateRelease[151] := BenchUut14.ActivateRelease;
   BenchCalls := BenchCalls + 1;
 152:
   BenchUut14.ManualMode := FALSE;
   BenchUut14.SingleStepMode := TRUE;
   BenchUut14.SingleCycleMode := FALSE;
   BenchUut14.ContinuousMode := FALSE;
   BenchUut14.EmergencyStop := TRUE;
   BenchUut14.Start := TRUE;
   BenchUut14.DownButton := FALSE;
   BenchUut14.UpButton := FALSE;
   BenchUut14.LeftButton := FALSE;
   BenchUut14.RightButton := FALSE;
   BenchUut14.GripButton := FALSE;
   BenchUut14.ReleaseButton := FALSE;
   BenchUut14.DownLimitSwitch := FALSE;
   BenchUut14.UpLimitSwitch := FALSE;
   BenchUut14.LeftLimitSwitch := FALSE;
   BenchUut14.RightLimitSwitch := FALSE;
   BenchUut14.GripLimitSwitch := FALSE;
   BenchUut14.ReleaseLimitSwitch := FALSE;
   TraceIn_ManualMode[152] := BenchUut14.ManualMode;
   TraceIn_SingleStepMode[152] := BenchUut14.SingleStepMode;
   TraceIn_SingleCycleMode[152] := BenchUut14.SingleCycleMode;
   TraceIn_ContinuousMode[152] := BenchUut14.ContinuousMode;
   TraceIn_EmergencyStop[152] := BenchUut14.EmergencyStop;
   TraceIn_Start[152] := BenchUut14.Start;
   TraceIn_DownButton[152] := BenchUut14.DownButton;
   TraceIn_UpButton[152] := BenchUut14.UpButton;
   TraceIn_LeftButton[152] := BenchUut14.LeftButton;
   TraceIn_RightButton[152] := BenchUut14.RightButton;
   TraceIn_GripButton[152] := BenchUut14.GripButton;
   TraceIn_ReleaseButton[152] := BenchUut14.ReleaseButton;
   TraceIn_DownLimitSwitch[152] := BenchUut14.DownLimitSwitch;
   TraceIn_UpLimitSwitch[152] := BenchUut14.UpLimitSwitch;
   TraceIn_LeftLimitSwitch[152] := BenchUut14.LeftLimitSwitch;
   TraceIn_RightLimitSwitch[152] := BenchUut14.RightLimitSwitch;
   TraceIn_GripLimitSwitch[152] := BenchUut14.GripLimitSwitch;
   TraceIn_ReleaseLimitSwitch[152] := BenchUut14.ReleaseLimitSwitch;
   BenchUut14();
   TraceOut_MoveDown[152] := BenchUut14.MoveDown;
   TraceOut_MoveUp[152] := BenchUut14.MoveUp;
   TraceOut_MoveLeft[152] := BenchUut14.MoveLeft;
   TraceOut_MoveRight[152] := BenchUut14.MoveRight;
   TraceOut_ActivateGrip[152] := BenchUut14.ActivateGrip;
   TraceOut_ActivateRelease[152] := BenchUut14.ActivateRelease;
   BenchCalls := BenchCalls + 1;
 153:
   BenchUut14.ManualMode := FALSE;
   BenchUut14.SingleStepMode := TRUE;
   BenchUut14.SingleCycleMode := FALSE;
   BenchUut14.ContinuousMode := FALSE;
   BenchUut14.EmergencyStop := TRUE;
   BenchUut14.Start := FALSE;
   BenchUut14.DownButton := FALSE;
   BenchUut14.UpButton := FALSE;
   BenchUut14.LeftButton := FALSE;
   BenchUut14.RightButton := FALSE;
   BenchUut14.GripButton := FALSE;
   BenchUut14.ReleaseButton := FALSE;
   BenchUut14.DownLimitSwitch := FALSE;
   BenchUut14.UpLimitSwitch := FALSE;
   BenchUut14.LeftLimitSwitch := FALSE;
   BenchUut14.RightLimitSwitch := FALSE;
   BenchUut14.GripLimitSwitch := FALSE;
   BenchUut14.ReleaseLimitSwitch := FALSE;
   TraceIn_ManualMode[153] := BenchUut14.ManualMode;
   TraceIn_SingleStepMode[153] := BenchUut14.SingleStepMode;
   TraceIn_SingleCycleMode[153] := BenchUut14.SingleCycleMode;
   TraceIn_ContinuousMode[153] := BenchUut14.ContinuousMode;
   TraceIn_EmergencyStop[153] := BenchUut14.EmergencyStop;
   TraceIn_Start[153] := BenchUut14.Start;
   TraceIn_DownButton[153] := BenchUut14.DownButton;
   TraceIn_UpButton[153] := BenchUut14.UpButton;
   TraceIn_LeftButton[153] := BenchUut14.LeftButton;
   TraceIn_RightButton[153] := BenchUut14.RightButton;
   TraceIn_GripButton[153] := BenchUut14.GripButton;
   TraceIn_ReleaseButton[153] := BenchUut14.ReleaseButton;
   TraceIn_DownLimitSwitch[153] := BenchUut14.DownLimitSwitch;
   TraceIn_UpLimitSwitch[153] := BenchUut14.UpLimitSwitch;
   TraceIn_LeftLimitSwitch[153] := BenchUut14.LeftLimitSwitch;
   TraceIn_RightLimitSwitch[153] := BenchUut14.RightLimitSwitch;
   TraceIn_GripLimitSwitch[153] := BenchUut14.GripLimitSwitch;
   TraceIn_ReleaseLimitSwitch[153] := BenchUut14.ReleaseLimitSwitch;
   BenchUut14();
   TraceOut_MoveDown[153] := BenchUut14.MoveDown;
   TraceOut_MoveUp[153] := BenchUut14.MoveUp;
   TraceOut_MoveLeft[153] := BenchUut14.MoveLeft;
   TraceOut_MoveRight[153] := BenchUut14.MoveRight;
   TraceOut_ActivateGrip[153] := BenchUut14.ActivateGrip;
   TraceOut_ActivateRelease[153] := BenchUut14.ActivateRelease;
   BenchCalls := BenchCalls + 1;
 154:
   BenchUut14.ManualMode := FALSE;
   BenchUut14.SingleStepMode := TRUE;
   BenchUut14.SingleCycleMode := FALSE;
   BenchUut14.ContinuousMode := FALSE;
   BenchUut14.EmergencyStop := TRUE;
   BenchUut14.Start := FALSE;
   BenchUut14.DownButton := FALSE;
   BenchUut14.UpButton := FALSE;
   BenchUut14.LeftButton := FALSE;
   BenchUut14.RightButton := FALSE;
   BenchUut14.GripButton := FALSE;
   BenchUut14.ReleaseButton := FALSE;
   BenchUut14.DownLimitSwitch := FALSE;
   BenchUut14.UpLimitSwitch := FALSE;
   BenchUut14.LeftLimitSwitch := FALSE;
   BenchUut14.RightLimitSwitch := FALSE;
   BenchUut14.GripLimitSwitch := FALSE;
   BenchUut14.ReleaseLimitSwitch := FALSE;
   TraceIn_ManualMode[154] := BenchUut14.ManualMode;
   TraceIn_SingleStepMode[154] := BenchUut14.SingleStepMode;
   TraceIn_SingleCycleMode[154] := BenchUut14.SingleCycleMode;
   TraceIn_ContinuousMode[154] := BenchUut14.ContinuousMode;
   TraceIn_EmergencyStop[154] := BenchUut14.EmergencyStop;
   TraceIn_Start[154] := BenchUut14.Start;
   TraceIn_DownButton[154] := BenchUut14.DownButton;
   TraceIn_UpButton[154] := BenchUut14.UpButton;
   TraceIn_LeftButton[154] := BenchUut14.LeftButton;
   TraceIn_RightButton[154] := BenchUut14.RightButton;
   TraceIn_GripButton[154] := BenchUut14.GripButton;
   TraceIn_ReleaseButton[154] := BenchUut14.ReleaseButton;
   TraceIn_DownLimitSwitch[154] := BenchUut14.DownLimitSwitch;
   TraceIn_UpLimitSwitch[154] := BenchUut14.UpLimitSwitch;
   TraceIn_LeftLimitSwitch[154] := BenchUut14.LeftLimitSwitch;
   TraceIn_RightLimitSwitch[154] := BenchUut14.RightLimitSwitch;
   TraceIn_GripLimitSwitch[154] := BenchUut14.GripLimitSwitch;
   TraceIn_ReleaseLimitSwitch[154] := BenchUut14.ReleaseLimitSwitch;
   BenchUut14();
   TraceOut_MoveDown[154] := BenchUut14.MoveDown;
   TraceOut_MoveUp[154] := BenchUut14.MoveUp;
   TraceOut_MoveLeft[154] := BenchUut14.MoveLeft;
   TraceOut_MoveRight[154] := BenchUut14.MoveRight;
   TraceOut_ActivateGrip[154] := BenchUut14.ActivateGrip;
   TraceOut_ActivateRelease[154] := BenchUut14.ActivateRelease;
   BenchCalls := BenchCalls + 1;
 155:
   BenchUut14.ManualMode := FALSE;
   BenchUut14.SingleStepMode := TRUE;
   BenchUut14.SingleCycleMode := FALSE;
   BenchUut14.ContinuousMode := FALSE;
   BenchUut14.EmergencyStop := TRUE;
   BenchUut14.Start := FALSE;
   BenchUut14.DownButton := FALSE;
   BenchUut14.UpButton := FALSE;
   BenchUut14.LeftButton := FALSE;
   BenchUut14.RightButton := FALSE;
   BenchUut14.GripButton := FALSE;
   BenchUut14.ReleaseButton := FALSE;
   BenchUut14.DownLimitSwitch := FALSE;
   BenchUut14.UpLimitSwitch := TRUE;
   BenchUut14.LeftLimitSwitch := FALSE;
   BenchUut14.RightLimitSwitch := FALSE;
   BenchUut14.GripLimitSwitch := FALSE;
   BenchUut14.ReleaseLimitSwitch := FALSE;
   TraceIn_ManualMode[155] := BenchUut14.ManualMode;
   TraceIn_SingleStepMode[155] := BenchUut14.SingleStepMode;
   TraceIn_SingleCycleMode[155] := BenchUut14.SingleCycleMode;
   TraceIn_ContinuousMode[155] := BenchUut14.ContinuousMode;
   TraceIn_EmergencyStop[155] := BenchUut14.EmergencyStop;
   TraceIn_Start[155] := BenchUut14.Start;
   TraceIn_DownButton[155] := BenchUut14.DownButton;
   TraceIn_UpButton[155] := BenchUut14.UpButton;
   TraceIn_LeftButton[155] := BenchUut14.LeftButton;
   TraceIn_RightButton[155] := BenchUut14.RightButton;
   TraceIn_GripButton[155] := BenchUut14.GripButton;
   TraceIn_ReleaseButton[155] := BenchUut14.ReleaseButton;
   TraceIn_DownLimitSwitch[155] := BenchUut14.DownLimitSwitch;
   TraceIn_UpLimitSwitch[155] := BenchUut14.UpLimitSwitch;
   TraceIn_LeftLimitSwitch[155] := BenchUut14.LeftLimitSwitch;
   TraceIn_RightLimitSwitch[155] := BenchUut14.RightLimitSwitch;
   TraceIn_GripLimitSwitch[155] := BenchUut14.GripLimitSwitch;
   TraceIn_ReleaseLimitSwitch[155] := BenchUut14.ReleaseLimitSwitch;
   BenchUut14();
   TraceOut_MoveDown[155] := BenchUut14.MoveDown;
   TraceOut_MoveUp[155] := BenchUut14.MoveUp;
   TraceOut_MoveLeft[155] := BenchUut14.MoveLeft;
   TraceOut_MoveRight[155] := BenchUut14.MoveRight;
   TraceOut_ActivateGrip[155] := BenchUut14.ActivateGrip;
   TraceOut_ActivateRelease[155] := BenchUut14.ActivateRelease;
   BenchCalls := BenchCalls + 1;
 156:
   BenchUut14.ManualMode := FALSE;
   BenchUut14.SingleStepMode := TRUE;
   BenchUut14.SingleCycleMode := FALSE;
   BenchUut14.ContinuousMode := FALSE;
   BenchUut14.EmergencyStop := TRUE;
   BenchUut14.Start := TRUE;
   BenchUut14.DownButton := FALSE;
   BenchUut14.UpButton := FALSE;
   BenchUut14.LeftButton := FALSE;
   BenchUut14.RightButton := FALSE;
   BenchUut14.GripButton := FALSE;
   BenchUut14.ReleaseButton := FALSE;
   BenchUut14.DownLimitSwitch := FALSE;
   BenchUut14.UpLimitSwitch := FALSE;
   BenchUut14.LeftLimitSwitch := FALSE;
   BenchUut14.RightLimitSwitch := FALSE;
   BenchUut14.GripLimitSwitch := FALSE;
   BenchUut14.ReleaseLimitSwitch := FALSE;
   TraceIn_ManualMode[156] := BenchUut14.ManualMode;
   TraceIn_SingleStepMode[156] := BenchUut14.SingleStepMode;
   TraceIn_SingleCycleMode[156] := BenchUut14.SingleCycleMode;
   TraceIn_ContinuousMode[156] := BenchUut14.ContinuousMode;
   TraceIn_EmergencyStop[156] := BenchUut14.EmergencyStop;
   TraceIn_Start[156] := BenchUut14.Start;
   TraceIn_DownButton[156] := BenchUut14.DownButton;
   TraceIn_UpButton[156] := BenchUut14.UpButton;
   TraceIn_LeftButton[156] := BenchUut14.LeftButton;
   TraceIn_RightButton[156] := BenchUut14.RightButton;
   TraceIn_GripButton[156] := BenchUut14.GripButton;
   TraceIn_ReleaseButton[156] := BenchUut14.ReleaseButton;
   TraceIn_DownLimitSwitch[156] := BenchUut14.DownLimitSwitch;
   TraceIn_UpLimitSwitch[156] := BenchUut14.UpLimitSwitch;
   TraceIn_LeftLimitSwitch[156] := BenchUut14.LeftLimitSwitch;
   TraceIn_RightLimitSwitch[156] := BenchUut14.RightLimitSwitch;
   TraceIn_GripLimitSwitch[156] := BenchUut14.GripLimitSwitch;
   TraceIn_ReleaseLimitSwitch[156] := BenchUut14.ReleaseLimitSwitch;
   BenchUut14();
   TraceOut_MoveDown[156] := BenchUut14.MoveDown;
   TraceOut_MoveUp[156] := BenchUut14.MoveUp;
   TraceOut_MoveLeft[156] := BenchUut14.MoveLeft;
   TraceOut_MoveRight[156] := BenchUut14.MoveRight;
   TraceOut_ActivateGrip[156] := BenchUut14.ActivateGrip;
   TraceOut_ActivateRelease[156] := BenchUut14.ActivateRelease;
   BenchCalls := BenchCalls + 1;
 157:
   BenchUut14.ManualMode := FALSE;
   BenchUut14.SingleStepMode := TRUE;
   BenchUut14.SingleCycleMode := FALSE;
   BenchUut14.ContinuousMode := FALSE;
   BenchUut14.EmergencyStop := TRUE;
   BenchUut14.Start := FALSE;
   BenchUut14.DownButton := FALSE;
   BenchUut14.UpButton := FALSE;
   BenchUut14.LeftButton := FALSE;
   BenchUut14.RightButton := FALSE;
   BenchUut14.GripButton := FALSE;
   BenchUut14.ReleaseButton := FALSE;
   BenchUut14.DownLimitSwitch := FALSE;
   BenchUut14.UpLimitSwitch := FALSE;
   BenchUut14.LeftLimitSwitch := FALSE;
   BenchUut14.RightLimitSwitch := FALSE;
   BenchUut14.GripLimitSwitch := FALSE;
   BenchUut14.ReleaseLimitSwitch := FALSE;
   TraceIn_ManualMode[157] := BenchUut14.ManualMode;
   TraceIn_SingleStepMode[157] := BenchUut14.SingleStepMode;
   TraceIn_SingleCycleMode[157] := BenchUut14.SingleCycleMode;
   TraceIn_ContinuousMode[157] := BenchUut14.ContinuousMode;
   TraceIn_EmergencyStop[157] := BenchUut14.EmergencyStop;
   TraceIn_Start[157] := BenchUut14.Start;
   TraceIn_DownButton[157] := BenchUut14.DownButton;
   TraceIn_UpButton[157] := BenchUut14.UpButton;
   TraceIn_LeftButton[157] := BenchUut14.LeftButton;
   TraceIn_RightButton[157] := BenchUut14.RightButton;
   TraceIn_GripButton[157] := BenchUut14.GripButton;
   TraceIn_ReleaseButton[157] := BenchUut14.ReleaseButton;
   TraceIn_DownLimitSwitch[157] := BenchUut14.DownLimitSwitch;
   TraceIn_UpLimitSwitch[157] := BenchUut14.UpLimitSwitch;
   TraceIn_LeftLimitSwitch[157] := BenchUut14.LeftLimitSwitch;
   TraceIn_RightLimitSwitch[157] := BenchUut14.RightLimitSwitch;
   TraceIn_GripLimitSwitch[157] := BenchUut14.GripLimitSwitch;
   TraceIn_ReleaseLimitSwitch[157] := BenchUut14.ReleaseLimitSwitch;
   BenchUut14();
   TraceOut_MoveDown[157] := BenchUut14.MoveDown;
   TraceOut_MoveUp[157] := BenchUut14.MoveUp;
   TraceOut_MoveLeft[157] := BenchUut14.MoveLeft;
   TraceOut_MoveRight[157] := BenchUut14.MoveRight;
   TraceOut_ActivateGrip[157] := BenchUut14.ActivateGrip;
   TraceOut_ActivateRelease[157] := BenchUut14.ActivateRelease;
   BenchCalls := BenchCalls + 1;
 158:
   BenchUut14.ManualMode := FALSE;
   BenchUut14.SingleStepMode := TRUE;
   BenchUut14.SingleCycleMode := FALSE;
   BenchUut14.ContinuousMode := FALSE;
   BenchUut14.EmergencyStop := TRUE;
   BenchUut14.Start := FALSE;
   BenchUut14.DownButton := FALSE;
   BenchUut14.UpButton := FALSE;
   BenchUut14.LeftButton := FALSE;
   BenchUut14.RightButton := FALSE;
   BenchUut14.GripButton := FALSE;
   BenchUut14.ReleaseButton := FALSE;
   BenchUut14.DownLimitSwitch := FALSE;
   BenchUut14.UpLimitSwitch := FALSE;
   BenchUut14.LeftLimitSwitch := FALSE;
   BenchUut14.RightLimitSwitch := FALSE;
   BenchUut14.GripLimitSwitch := FALSE;
   BenchUut14.ReleaseLimitSwitch := FALSE;
   TraceIn_ManualMode[158] := BenchUut14.ManualMode;
   TraceIn_SingleStepMode[158] := BenchUut14.SingleStepMode;
   TraceIn_SingleCycleMode[158] := BenchUut14.SingleCycleMode;
   TraceIn_ContinuousMode[158] := BenchUut14.ContinuousMode;
   TraceIn_EmergencyStop[158] := BenchUut14.EmergencyStop;
   TraceIn_Start[158] := BenchUut14.Start;
   TraceIn_DownButton[158] := BenchUut14.DownButton;
   TraceIn_UpButton[158] := BenchUut14.UpButton;
   TraceIn_LeftButton[158] := BenchUut14.LeftButton;
   TraceIn_RightButton[158] := BenchUut14.RightButton;
   TraceIn_GripButton[158] := BenchUut14.GripButton;
   TraceIn_ReleaseButton[158] := BenchUut14.ReleaseButton;
   TraceIn_DownLimitSwitch[158] := BenchUut14.DownLimitSwitch;
   TraceIn_UpLimitSwitch[158] := BenchUut14.UpLimitSwitch;
   TraceIn_LeftLimitSwitch[158] := BenchUut14.LeftLimitSwitch;
   TraceIn_RightLimitSwitch[158] := BenchUut14.RightLimitSwitch;
   TraceIn_GripLimitSwitch[158] := BenchUut14.GripLimitSwitch;
   TraceIn_ReleaseLimitSwitch[158] := BenchUut14.ReleaseLimitSwitch;
   BenchUut14();
   TraceOut_MoveDown[158] := BenchUut14.MoveDown;
   TraceOut_MoveUp[158] := BenchUut14.MoveUp;
   TraceOut_MoveLeft[158] := BenchUut14.MoveLeft;
   TraceOut_MoveRight[158] := BenchUut14.MoveRight;
   TraceOut_ActivateGrip[158] := BenchUut14.ActivateGrip;
   TraceOut_ActivateRelease[158] := BenchUut14.ActivateRelease;
   BenchCalls := BenchCalls + 1;
 159:
   BenchUut14.ManualMode := FALSE;
   BenchUut14.SingleStepMode := TRUE;
   BenchUut14.SingleCycleMode := FALSE;
   BenchUut14.ContinuousMode := FALSE;
   BenchUut14.EmergencyStop := TRUE;
   BenchUut14.Start := FALSE;
   BenchUut14.DownButton := FALSE;
   BenchUut14.UpButton := FALSE;
   BenchUut14.LeftButton := FALSE;
   BenchUut14.RightButton := FALSE;
   BenchUut14.GripButton := FALSE;
   BenchUut14.ReleaseButton := FALSE;
   BenchUut14.DownLimitSwitch := FALSE;
   BenchUut14.UpLimitSwitch := FALSE;
   BenchUut14.LeftLimitSwitch := FALSE;
   BenchUut14.RightLimitSwitch := TRUE;
   BenchUut14.GripLimitSwitch := FALSE;
   BenchUut14.ReleaseLimitSwitch := FALSE;
   TraceIn_ManualMode[159] := BenchUut14.ManualMode;
   TraceIn_SingleStepMode[159] := BenchUut14.SingleStepMode;
   TraceIn_SingleCycleMode[159] := BenchUut14.SingleCycleMode;
   TraceIn_ContinuousMode[159] := BenchUut14.ContinuousMode;
   TraceIn_EmergencyStop[159] := BenchUut14.EmergencyStop;
   TraceIn_Start[159] := BenchUut14.Start;
   TraceIn_DownButton[159] := BenchUut14.DownButton;
   TraceIn_UpButton[159] := BenchUut14.UpButton;
   TraceIn_LeftButton[159] := BenchUut14.LeftButton;
   TraceIn_RightButton[159] := BenchUut14.RightButton;
   TraceIn_GripButton[159] := BenchUut14.GripButton;
   TraceIn_ReleaseButton[159] := BenchUut14.ReleaseButton;
   TraceIn_DownLimitSwitch[159] := BenchUut14.DownLimitSwitch;
   TraceIn_UpLimitSwitch[159] := BenchUut14.UpLimitSwitch;
   TraceIn_LeftLimitSwitch[159] := BenchUut14.LeftLimitSwitch;
   TraceIn_RightLimitSwitch[159] := BenchUut14.RightLimitSwitch;
   TraceIn_GripLimitSwitch[159] := BenchUut14.GripLimitSwitch;
   TraceIn_ReleaseLimitSwitch[159] := BenchUut14.ReleaseLimitSwitch;
   BenchUut14();
   TraceOut_MoveDown[159] := BenchUut14.MoveDown;
   TraceOut_MoveUp[159] := BenchUut14.MoveUp;
   TraceOut_MoveLeft[159] := BenchUut14.MoveLeft;
   TraceOut_MoveRight[159] := BenchUut14.MoveRight;
   TraceOut_ActivateGrip[159] := BenchUut14.ActivateGrip;
   TraceOut_ActivateRelease[159] := BenchUut14.ActivateRelease;
   BenchCalls := BenchCalls + 1;
 160:
   BenchUut14.ManualMode := FALSE;
   BenchUut14.SingleStepMode := TRUE;
   BenchUut14.SingleCycleMode := FALSE;
   BenchUut14.ContinuousMode := FALSE;
   BenchUut14.EmergencyStop := TRUE;
   BenchUut14.Start := TRUE;
   BenchUut14.DownButton := FALSE;
   BenchUut14.UpButton := FALSE;
   BenchUut14.LeftButton := FALSE;
   BenchUut14.RightButton := FALSE;
   BenchUut14.GripButton := FALSE;
   BenchUut14.ReleaseButton := FALSE;
   BenchUut14.DownLimitSwitch := FALSE;
   BenchUut14.UpLimitSwitch := FALSE;
   BenchUut14.LeftLimitSwitch := FALSE;
   BenchUut14.RightLimitSwitch := FALSE;
   BenchUut14.GripLimitSwitch := FALSE;
   BenchUut14.ReleaseLimitSwitch := FALSE;
   TraceIn_ManualMode[160] := BenchUut14.ManualMode;
   TraceIn_SingleStepMode[160] := BenchUut14.SingleStepMode;
   TraceIn_SingleCycleMode[160] := BenchUut14.SingleCycleMode;
   TraceIn_ContinuousMode[160] := BenchUut14.ContinuousMode;
   TraceIn_EmergencyStop[160] := BenchUut14.EmergencyStop;
   TraceIn_Start[160] := BenchUut14.Start;
   TraceIn_DownButton[160] := BenchUut14.DownButton;
   TraceIn_UpButton[160] := BenchUut14.UpButton;
   TraceIn_LeftButton[160] := BenchUut14.LeftButton;
   TraceIn_RightButton[160] := BenchUut14.RightButton;
   TraceIn_GripButton[160] := BenchUut14.GripButton;
   TraceIn_ReleaseButton[160] := BenchUut14.ReleaseButton;
   TraceIn_DownLimitSwitch[160] := BenchUut14.DownLimitSwitch;
   TraceIn_UpLimitSwitch[160] := BenchUut14.UpLimitSwitch;
   TraceIn_LeftLimitSwitch[160] := BenchUut14.LeftLimitSwitch;
   TraceIn_RightLimitSwitch[160] := BenchUut14.RightLimitSwitch;
   TraceIn_GripLimitSwitch[160] := BenchUut14.GripLimitSwitch;
   TraceIn_ReleaseLimitSwitch[160] := BenchUut14.ReleaseLimitSwitch;
   BenchUut14();
   TraceOut_MoveDown[160] := BenchUut14.MoveDown;
   TraceOut_MoveUp[160] := BenchUut14.MoveUp;
   TraceOut_MoveLeft[160] := BenchUut14.MoveLeft;
   TraceOut_MoveRight[160] := BenchUut14.MoveRight;
   TraceOut_ActivateGrip[160] := BenchUut14.ActivateGrip;
   TraceOut_ActivateRelease[160] := BenchUut14.ActivateRelease;
   BenchCalls := BenchCalls + 1;
 161:
   BenchUut14.ManualMode := FALSE;
   BenchUut14.SingleStepMode := TRUE;
   BenchUut14.SingleCycleMode := FALSE;
   BenchUut14.ContinuousMode := FALSE;
   BenchUut14.EmergencyStop := TRUE;
   BenchUut14.Start := FALSE;
   BenchUut14.DownButton := FALSE;
   BenchUut14.UpButton := FALSE;
   BenchUut14.LeftButton := FALSE;
   BenchUut14.RightButton := FALSE;
   BenchUut14.GripButton := FALSE;
   BenchUut14.ReleaseButton := FALSE;
   BenchUut14.DownLimitSwitch := FALSE;
   BenchUut14.UpLimitSwitch := FALSE;
   BenchUut14.LeftLimitSwitch := FALSE;
   BenchUut14.RightLimitSwitch := FALSE;
   BenchUut14.GripLimitSwitch := FALSE;
   BenchUut14.ReleaseLimitSwitch := FALSE;
   TraceIn_ManualMode[161] := BenchUut14.ManualMode;
   TraceIn_SingleStepMode[161] := BenchUut14.SingleStepMode;
   TraceIn_SingleCycleMode[161] := BenchUut14.SingleCycleMode;
   TraceIn_ContinuousMode[161] := BenchUut14.ContinuousMode;
   TraceIn_EmergencyStop[161] := BenchUut14.EmergencyStop;
   TraceIn_Start[161] := BenchUut14.Start;
   TraceIn_DownButton[161] := BenchUut14.DownButton;
   TraceIn_UpButton[161] := BenchUut14.UpButton;
   TraceIn_LeftButton[161] := BenchUut14.LeftButton;
   TraceIn_RightButton[161] := BenchUut14.RightButton;
   TraceIn_GripButton[161] := BenchUut14.GripButton;
   TraceIn_ReleaseButton[161] := BenchUut14.ReleaseButton;
   TraceIn_DownLimitSwitch[161] := BenchUut14.DownLimitSwitch;
   TraceIn_UpLimitSwitch[161] := BenchUut14.UpLimitSwitch;
   TraceIn_LeftLimitSwitch[161] := BenchUut14.LeftLimitSwitch;
   TraceIn_RightLimitSwitch[161] := BenchUut14.RightLimitSwitch;
   TraceIn_GripLimitSwitch[161] := BenchUut14.GripLimitSwitch;
   TraceIn_ReleaseLimitSwitch[161] := BenchUut14.ReleaseLimitSwitch;
   BenchUut14();
   TraceOut_MoveDown[161] := BenchUut14.MoveDown;
   TraceOut_MoveUp[161] := BenchUut14.MoveUp;
   TraceOut_MoveLeft[161] := BenchUut14.MoveLeft;
   TraceOut_MoveRight[161] := BenchUut14.MoveRight;
   TraceOut_ActivateGrip[161] := BenchUut14.ActivateGrip;
   TraceOut_ActivateRelease[161] := BenchUut14.ActivateRelease;
   BenchCalls := BenchCalls + 1;
 162:
   BenchUut14.ManualMode := FALSE;
   BenchUut14.SingleStepMode := TRUE;
   BenchUut14.SingleCycleMode := FALSE;
   BenchUut14.ContinuousMode := FALSE;
   BenchUut14.EmergencyStop := TRUE;
   BenchUut14.Start := FALSE;
   BenchUut14.DownButton := FALSE;
   BenchUut14.UpButton := FALSE;
   BenchUut14.LeftButton := FALSE;
   BenchUut14.RightButton := FALSE;
   BenchUut14.GripButton := FALSE;
   BenchUut14.ReleaseButton := FALSE;
   BenchUut14.DownLimitSwitch := FALSE;
   BenchUut14.UpLimitSwitch := FALSE;
   BenchUut14.LeftLimitSwitch := FALSE;
   BenchUut14.RightLimitSwitch := FALSE;
   BenchUut14.GripLimitSwitch := FALSE;
   BenchUut14.ReleaseLimitSwitch := FALSE;
   TraceIn_ManualMode[162] := BenchUut14.ManualMode;
   TraceIn_SingleStepMode[162] := BenchUut14.SingleStepMode;
   TraceIn_SingleCycleMode[162] := BenchUut14.SingleCycleMode;
   TraceIn_ContinuousMode[162] := BenchUut14.ContinuousMode;
   TraceIn_EmergencyStop[162] := BenchUut14.EmergencyStop;
   TraceIn_Start[162] := BenchUut14.Start;
   TraceIn_DownButton[162] := BenchUut14.DownButton;
   TraceIn_UpButton[162] := BenchUut14.UpButton;
   TraceIn_LeftButton[162] := BenchUut14.LeftButton;
   TraceIn_RightButton[162] := BenchUut14.RightButton;
   TraceIn_GripButton[162] := BenchUut14.GripButton;
   TraceIn_ReleaseButton[162] := BenchUut14.ReleaseButton;
   TraceIn_DownLimitSwitch[162] := BenchUut14.DownLimitSwitch;
   TraceIn_UpLimitSwitch[162] := BenchUut14.UpLimitSwitch;
   TraceIn_LeftLimitSwitch[162] := BenchUut14.LeftLimitSwitch;
   TraceIn_RightLimitSwitch[162] := BenchUut14.RightLimitSwitch;
   TraceIn_GripLimitSwitch[162] := BenchUut14.GripLimitSwitch;
   TraceIn_ReleaseLimitSwitch[162] := BenchUut14.ReleaseLimitSwitch;
   BenchUut14();
   TraceOut_MoveDown[162] := BenchUut14.MoveDown;
   TraceOut_MoveUp[162] := BenchUut14.MoveUp;
   TraceOut_MoveLeft[162] := BenchUut14.MoveLeft;
   TraceOut_MoveRight[162] := BenchUut14.MoveRight;
   TraceOut_ActivateGrip[162] := BenchUut14.ActivateGrip;
   TraceOut_ActivateRelease[162] := BenchUut14.ActivateRelease;
   BenchCalls := BenchCalls + 1;
 163:
   BenchUut14.ManualMode := FALSE;
   BenchUut14.SingleStepMode := TRUE;
   BenchUut14.SingleCycleMode := FALSE;
   BenchUut14.ContinuousMode := FALSE;
   BenchUut14.EmergencyStop := TRUE;
   BenchUut14.Start := FALSE;
   BenchUut14.DownButton := FALSE;
   BenchUut14.UpButton := FALSE;
   BenchUut14.LeftButton := FALSE;
   BenchUut14.RightButton := FALSE;
   BenchUut14.GripButton := FALSE;
   BenchUut14.ReleaseButton := FALSE;
   BenchUut14.DownLimitSwitch := TRUE;
   BenchUut14.UpLimitSwitch := FALSE;
   BenchUut14.LeftLimitSwitch := FALSE;
   BenchUut14.RightLimitSwitch := FALSE;
   BenchUut14.GripLimitSwitch := FALSE;
   BenchUut14.ReleaseLimitSwitch := FALSE;
   TraceIn_ManualMode[163] := BenchUut14.ManualMode;
   TraceIn_SingleStepMode[163] := BenchUut14.SingleStepMode;
   TraceIn_SingleCycleMode[163] := BenchUut14.SingleCycleMode;
   TraceIn_ContinuousMode[163] := BenchUut14.ContinuousMode;
   TraceIn_EmergencyStop[163] := BenchUut14.EmergencyStop;
   TraceIn_Start[163] := BenchUut14.Start;
   TraceIn_DownButton[163] := BenchUut14.DownButton;
   TraceIn_UpButton[163] := BenchUut14.UpButton;
   TraceIn_LeftButton[163] := BenchUut14.LeftButton;
   TraceIn_RightButton[163] := BenchUut14.RightButton;
   TraceIn_GripButton[163] := BenchUut14.GripButton;
   TraceIn_ReleaseButton[163] := BenchUut14.ReleaseButton;
   TraceIn_DownLimitSwitch[163] := BenchUut14.DownLimitSwitch;
   TraceIn_UpLimitSwitch[163] := BenchUut14.UpLimitSwitch;
   TraceIn_LeftLimitSwitch[163] := BenchUut14.LeftLimitSwitch;
   TraceIn_RightLimitSwitch[163] := BenchUut14.RightLimitSwitch;
   TraceIn_GripLimitSwitch[163] := BenchUut14.GripLimitSwitch;
   TraceIn_ReleaseLimitSwitch[163] := BenchUut14.ReleaseLimitSwitch;
   BenchUut14();
   TraceOut_MoveDown[163] := BenchUut14.MoveDown;
   TraceOut_MoveUp[163] := BenchUut14.MoveUp;
   TraceOut_MoveLeft[163] := BenchUut14.MoveLeft;
   TraceOut_MoveRight[163] := BenchUut14.MoveRight;
   TraceOut_ActivateGrip[163] := BenchUut14.ActivateGrip;
   TraceOut_ActivateRelease[163] := BenchUut14.ActivateRelease;
   BenchCalls := BenchCalls + 1;
 164:
   BenchUut14.ManualMode := FALSE;
   BenchUut14.SingleStepMode := TRUE;
   BenchUut14.SingleCycleMode := FALSE;
   BenchUut14.ContinuousMode := FALSE;
   BenchUut14.EmergencyStop := TRUE;
   BenchUut14.Start := TRUE;
   BenchUut14.DownButton := FALSE;
   BenchUut14.UpButton := FALSE;
   BenchUut14.LeftButton := FALSE;
   BenchUut14.RightButton := FALSE;
   BenchUut14.GripButton := FALSE;
   BenchUut14.ReleaseButton := FALSE;
   BenchUut14.DownLimitSwitch := FALSE;
   BenchUut14.UpLimitSwitch := FALSE;
   BenchUut14.LeftLimitSwitch := FALSE;
   BenchUut14.RightLimitSwitch := FALSE;
   BenchUut14.GripLimitSwitch := FALSE;
   BenchUut14.ReleaseLimitSwitch := FALSE;
   TraceIn_ManualMode[164] := BenchUut14.ManualMode;
   TraceIn_SingleStepMode[164] := BenchUut14.SingleStepMode;
   TraceIn_SingleCycleMode[164] := BenchUut14.SingleCycleMode;
   TraceIn_ContinuousMode[164] := BenchUut14.ContinuousMode;
   TraceIn_EmergencyStop[164] := BenchUut14.EmergencyStop;
   TraceIn_Start[164] := BenchUut14.Start;
   TraceIn_DownButton[164] := BenchUut14.DownButton;
   TraceIn_UpButton[164] := BenchUut14.UpButton;
   TraceIn_LeftButton[164] := BenchUut14.LeftButton;
   TraceIn_RightButton[164] := BenchUut14.RightButton;
   TraceIn_GripButton[164] := BenchUut14.GripButton;
   TraceIn_ReleaseButton[164] := BenchUut14.ReleaseButton;
   TraceIn_DownLimitSwitch[164] := BenchUut14.DownLimitSwitch;
   TraceIn_UpLimitSwitch[164] := BenchUut14.UpLimitSwitch;
   TraceIn_LeftLimitSwitch[164] := BenchUut14.LeftLimitSwitch;
   TraceIn_RightLimitSwitch[164] := BenchUut14.RightLimitSwitch;
   TraceIn_GripLimitSwitch[164] := BenchUut14.GripLimitSwitch;
   TraceIn_ReleaseLimitSwitch[164] := BenchUut14.ReleaseLimitSwitch;
   BenchUut14();
   TraceOut_MoveDown[164] := BenchUut14.MoveDown;
   TraceOut_MoveUp[164] := BenchUut14.MoveUp;
   TraceOut_MoveLeft[164] := BenchUut14.MoveLeft;
   TraceOut_MoveRight[164] := BenchUut14.MoveRight;
   TraceOut_ActivateGrip[164] := BenchUut14.ActivateGrip;
   TraceOut_ActivateRelease[164] := BenchUut14.ActivateRelease;
   BenchCalls := BenchCalls + 1;
 165:
   BenchUut14.ManualMode := FALSE;
   BenchUut14.SingleStepMode := TRUE;
   BenchUut14.SingleCycleMode := FALSE;
   BenchUut14.ContinuousMode := FALSE;
   BenchUut14.EmergencyStop := TRUE;
   BenchUut14.Start := FALSE;
   BenchUut14.DownButton := FALSE;
   BenchUut14.UpButton := FALSE;
   BenchUut14.LeftButton := FALSE;
   BenchUut14.RightButton := FALSE;
   BenchUut14.GripButton := FALSE;
   BenchUut14.ReleaseButton := FALSE;
   BenchUut14.DownLimitSwitch := FALSE;
   BenchUut14.UpLimitSwitch := FALSE;
   BenchUut14.LeftLimitSwitch := FALSE;
   BenchUut14.RightLimitSwitch := FALSE;
   BenchUut14.GripLimitSwitch := FALSE;
   BenchUut14.ReleaseLimitSwitch := FALSE;
   TraceIn_ManualMode[165] := BenchUut14.ManualMode;
   TraceIn_SingleStepMode[165] := BenchUut14.SingleStepMode;
   TraceIn_SingleCycleMode[165] := BenchUut14.SingleCycleMode;
   TraceIn_ContinuousMode[165] := BenchUut14.ContinuousMode;
   TraceIn_EmergencyStop[165] := BenchUut14.EmergencyStop;
   TraceIn_Start[165] := BenchUut14.Start;
   TraceIn_DownButton[165] := BenchUut14.DownButton;
   TraceIn_UpButton[165] := BenchUut14.UpButton;
   TraceIn_LeftButton[165] := BenchUut14.LeftButton;
   TraceIn_RightButton[165] := BenchUut14.RightButton;
   TraceIn_GripButton[165] := BenchUut14.GripButton;
   TraceIn_ReleaseButton[165] := BenchUut14.ReleaseButton;
   TraceIn_DownLimitSwitch[165] := BenchUut14.DownLimitSwitch;
   TraceIn_UpLimitSwitch[165] := BenchUut14.UpLimitSwitch;
   TraceIn_LeftLimitSwitch[165] := BenchUut14.LeftLimitSwitch;
   TraceIn_RightLimitSwitch[165] := BenchUut14.RightLimitSwitch;
   TraceIn_GripLimitSwitch[165] := BenchUut14.GripLimitSwitch;
   TraceIn_ReleaseLimitSwitch[165] := BenchUut14.ReleaseLimitSwitch;
   BenchUut14();
   TraceOut_MoveDown[165] := BenchUut14.MoveDown;
   TraceOut_MoveUp[165] := BenchUut14.MoveUp;
   TraceOut_MoveLeft[165] := BenchUut14.MoveLeft;
   TraceOut_MoveRight[165] := BenchUut14.MoveRight;
   TraceOut_ActivateGrip[165] := BenchUut14.ActivateGrip;
   TraceOut_ActivateRelease[165] := BenchUut14.ActivateRelease;
   BenchCalls := BenchCalls + 1;
 166:
   BenchUut14.ManualMode := FALSE;
   BenchUut14.SingleStepMode := TRUE;
   BenchUut14.SingleCycleMode := FALSE;
   BenchUut14.ContinuousMode := FALSE;
   BenchUut14.EmergencyStop := TRUE;
   BenchUut14.Start := FALSE;
   BenchUut14.DownButton := FALSE;
   BenchUut14.UpButton := FALSE;
   BenchUut14.LeftButton := FALSE;
   BenchUut14.RightButton := FALSE;
   BenchUut14.GripButton := FALSE;
   BenchUut14.ReleaseButton := FALSE;
   BenchUut14.DownLimitSwitch := FALSE;
   BenchUut14.UpLimitSwitch := FALSE;
   BenchUut14.LeftLimitSwitch := FALSE;
   BenchUut14.RightLimitSwitch := FALSE;
   BenchUut14.GripLimitSwitch := FALSE;
   BenchUut14.ReleaseLimitSwitch := FALSE;
   TraceIn_ManualMode[166] := BenchUut14.ManualMode;
   TraceIn_SingleStepMode[166] := BenchUut14.SingleStepMode;
   TraceIn_SingleCycleMode[166] := BenchUut14.SingleCycleMode;
   TraceIn_ContinuousMode[166] := BenchUut14.ContinuousMode;
   TraceIn_EmergencyStop[166] := BenchUut14.EmergencyStop;
   TraceIn_Start[166] := BenchUut14.Start;
   TraceIn_DownButton[166] := BenchUut14.DownButton;
   TraceIn_UpButton[166] := BenchUut14.UpButton;
   TraceIn_LeftButton[166] := BenchUut14.LeftButton;
   TraceIn_RightButton[166] := BenchUut14.RightButton;
   TraceIn_GripButton[166] := BenchUut14.GripButton;
   TraceIn_ReleaseButton[166] := BenchUut14.ReleaseButton;
   TraceIn_DownLimitSwitch[166] := BenchUut14.DownLimitSwitch;
   TraceIn_UpLimitSwitch[166] := BenchUut14.UpLimitSwitch;
   TraceIn_LeftLimitSwitch[166] := BenchUut14.LeftLimitSwitch;
   TraceIn_RightLimitSwitch[166] := BenchUut14.RightLimitSwitch;
   TraceIn_GripLimitSwitch[166] := BenchUut14.GripLimitSwitch;
   TraceIn_ReleaseLimitSwitch[166] := BenchUut14.ReleaseLimitSwitch;
   BenchUut14();
   TraceOut_MoveDown[166] := BenchUut14.MoveDown;
   TraceOut_MoveUp[166] := BenchUut14.MoveUp;
   TraceOut_MoveLeft[166] := BenchUut14.MoveLeft;
   TraceOut_MoveRight[166] := BenchUut14.MoveRight;
   TraceOut_ActivateGrip[166] := BenchUut14.ActivateGrip;
   TraceOut_ActivateRelease[166] := BenchUut14.ActivateRelease;
   BenchCalls := BenchCalls + 1;
 167:
   BenchUut14.ManualMode := FALSE;
   BenchUut14.SingleStepMode := TRUE;
   BenchUut14.SingleCycleMode := FALSE;
   BenchUut14.ContinuousMode := FALSE;
   BenchUut14.EmergencyStop := TRUE;
   BenchUut14.Start := FALSE;
   BenchUut14.DownButton := FALSE;
   BenchUut14.UpButton := FALSE;
   BenchUut14.LeftButton := FALSE;
   BenchUut14.RightButton := FALSE;
   BenchUut14.GripButton := FALSE;
   BenchUut14.ReleaseButton := FALSE;
   BenchUut14.DownLimitSwitch := FALSE;
   BenchUut14.UpLimitSwitch := FALSE;
   BenchUut14.LeftLimitSwitch := FALSE;
   BenchUut14.RightLimitSwitch := FALSE;
   BenchUut14.GripLimitSwitch := FALSE;
   BenchUut14.ReleaseLimitSwitch := TRUE;
   TraceIn_ManualMode[167] := BenchUut14.ManualMode;
   TraceIn_SingleStepMode[167] := BenchUut14.SingleStepMode;
   TraceIn_SingleCycleMode[167] := BenchUut14.SingleCycleMode;
   TraceIn_ContinuousMode[167] := BenchUut14.ContinuousMode;
   TraceIn_EmergencyStop[167] := BenchUut14.EmergencyStop;
   TraceIn_Start[167] := BenchUut14.Start;
   TraceIn_DownButton[167] := BenchUut14.DownButton;
   TraceIn_UpButton[167] := BenchUut14.UpButton;
   TraceIn_LeftButton[167] := BenchUut14.LeftButton;
   TraceIn_RightButton[167] := BenchUut14.RightButton;
   TraceIn_GripButton[167] := BenchUut14.GripButton;
   TraceIn_ReleaseButton[167] := BenchUut14.ReleaseButton;
   TraceIn_DownLimitSwitch[167] := BenchUut14.DownLimitSwitch;
   TraceIn_UpLimitSwitch[167] := BenchUut14.UpLimitSwitch;
   TraceIn_LeftLimitSwitch[167] := BenchUut14.LeftLimitSwitch;
   TraceIn_RightLimitSwitch[167] := BenchUut14.RightLimitSwitch;
   TraceIn_GripLimitSwitch[167] := BenchUut14.GripLimitSwitch;
   TraceIn_ReleaseLimitSwitch[167] := BenchUut14.ReleaseLimitSwitch;
   BenchUut14();
   TraceOut_MoveDown[167] := BenchUut14.MoveDown;
   TraceOut_MoveUp[167] := BenchUut14.MoveUp;
   TraceOut_MoveLeft[167] := BenchUut14.MoveLeft;
   TraceOut_MoveRight[167] := BenchUut14.MoveRight;
   TraceOut_ActivateGrip[167] := BenchUut14.ActivateGrip;
   TraceOut_ActivateRelease[167] := BenchUut14.ActivateRelease;
   BenchCalls := BenchCalls + 1;
 168:
   BenchUut14.ManualMode := FALSE;
   BenchUut14.SingleStepMode := TRUE;
   BenchUut14.SingleCycleMode := FALSE;
   BenchUut14.ContinuousMode := FALSE;
   BenchUut14.EmergencyStop := TRUE;
   BenchUut14.Start := TRUE;
   BenchUut14.DownButton := FALSE;
   BenchUut14.UpButton := FALSE;
   BenchUut14.LeftButton := FALSE;
   BenchUut14.RightButton := FALSE;
   BenchUut14.GripButton := FALSE;
   BenchUut14.ReleaseButton := FALSE;
   BenchUut14.DownLimitSwitch := FALSE;
   BenchUut14.UpLimitSwitch := FALSE;
   BenchUut14.LeftLimitSwitch := FALSE;
   BenchUut14.RightLimitSwitch := FALSE;
   BenchUut14.GripLimitSwitch := FALSE;
   BenchUut14.ReleaseLimitSwitch := FALSE;
   TraceIn_ManualMode[168] := BenchUut14.ManualMode;
   TraceIn_SingleStepMode[168] := BenchUut14.SingleStepMode;
   TraceIn_SingleCycleMode[168] := BenchUut14.SingleCycleMode;
   TraceIn_ContinuousMode[168] := BenchUut14.ContinuousMode;
   TraceIn_EmergencyStop[168] := BenchUut14.EmergencyStop;
   TraceIn_Start[168] := BenchUut14.Start;
   TraceIn_DownButton[168] := BenchUut14.DownButton;
   TraceIn_UpButton[168] := BenchUut14.UpButton;
   TraceIn_LeftButton[168] := BenchUut14.LeftButton;
   TraceIn_RightButton[168] := BenchUut14.RightButton;
   TraceIn_GripButton[168] := BenchUut14.GripButton;
   TraceIn_ReleaseButton[168] := BenchUut14.ReleaseButton;
   TraceIn_DownLimitSwitch[168] := BenchUut14.DownLimitSwitch;
   TraceIn_UpLimitSwitch[168] := BenchUut14.UpLimitSwitch;
   TraceIn_LeftLimitSwitch[168] := BenchUut14.LeftLimitSwitch;
   TraceIn_RightLimitSwitch[168] := BenchUut14.RightLimitSwitch;
   TraceIn_GripLimitSwitch[168] := BenchUut14.GripLimitSwitch;
   TraceIn_ReleaseLimitSwitch[168] := BenchUut14.ReleaseLimitSwitch;
   BenchUut14();
   TraceOut_MoveDown[168] := BenchUut14.MoveDown;
   TraceOut_MoveUp[168] := BenchUut14.MoveUp;
   TraceOut_MoveLeft[168] := BenchUut14.MoveLeft;
   TraceOut_MoveRight[168] := BenchUut14.MoveRight;
   TraceOut_ActivateGrip[168] := BenchUut14.ActivateGrip;
   TraceOut_ActivateRelease[168] := BenchUut14.ActivateRelease;
   BenchCalls := BenchCalls + 1;
 169:
   BenchUut14.ManualMode := FALSE;
   BenchUut14.SingleStepMode := TRUE;
   BenchUut14.SingleCycleMode := FALSE;
   BenchUut14.ContinuousMode := FALSE;
   BenchUut14.EmergencyStop := TRUE;
   BenchUut14.Start := FALSE;
   BenchUut14.DownButton := FALSE;
   BenchUut14.UpButton := FALSE;
   BenchUut14.LeftButton := FALSE;
   BenchUut14.RightButton := FALSE;
   BenchUut14.GripButton := FALSE;
   BenchUut14.ReleaseButton := FALSE;
   BenchUut14.DownLimitSwitch := FALSE;
   BenchUut14.UpLimitSwitch := FALSE;
   BenchUut14.LeftLimitSwitch := FALSE;
   BenchUut14.RightLimitSwitch := FALSE;
   BenchUut14.GripLimitSwitch := FALSE;
   BenchUut14.ReleaseLimitSwitch := FALSE;
   TraceIn_ManualMode[169] := BenchUut14.ManualMode;
   TraceIn_SingleStepMode[169] := BenchUut14.SingleStepMode;
   TraceIn_SingleCycleMode[169] := BenchUut14.SingleCycleMode;
   TraceIn_ContinuousMode[169] := BenchUut14.ContinuousMode;
   TraceIn_EmergencyStop[169] := BenchUut14.EmergencyStop;
   TraceIn_Start[169] := BenchUut14.Start;
   TraceIn_DownButton[169] := BenchUut14.DownButton;
   TraceIn_UpButton[169] := BenchUut14.UpButton;
   TraceIn_LeftButton[169] := BenchUut14.LeftButton;
   TraceIn_RightButton[169] := BenchUut14.RightButton;
   TraceIn_GripButton[169] := BenchUut14.GripButton;
   TraceIn_ReleaseButton[169] := BenchUut14.ReleaseButton;
   TraceIn_DownLimitSwitch[169] := BenchUut14.DownLimitSwitch;
   TraceIn_UpLimitSwitch[169] := BenchUut14.UpLimitSwitch;
   TraceIn_LeftLimitSwitch[169] := BenchUut14.LeftLimitSwitch;
   TraceIn_RightLimitSwitch[169] := BenchUut14.RightLimitSwitch;
   TraceIn_GripLimitSwitch[169] := BenchUut14.GripLimitSwitch;
   TraceIn_ReleaseLimitSwitch[169] := BenchUut14.ReleaseLimitSwitch;
   BenchUut14();
   TraceOut_MoveDown[169] := BenchUut14.MoveDown;
   TraceOut_MoveUp[169] := BenchUut14.MoveUp;
   TraceOut_MoveLeft[169] := BenchUut14.MoveLeft;
   TraceOut_MoveRight[169] := BenchUut14.MoveRight;
   TraceOut_ActivateGrip[169] := BenchUut14.ActivateGrip;
   TraceOut_ActivateRelease[169] := BenchUut14.ActivateRelease;
   BenchCalls := BenchCalls + 1;
 170:
   BenchUut14.ManualMode := FALSE;
   BenchUut14.SingleStepMode := TRUE;
   BenchUut14.SingleCycleMode := FALSE;
   BenchUut14.ContinuousMode := FALSE;
   BenchUut14.EmergencyStop := TRUE;
   BenchUut14.Start := FALSE;
   BenchUut14.DownButton := FALSE;
   BenchUut14.UpButton := FALSE;
   BenchUut14.LeftButton := FALSE;
   BenchUut14.RightButton := FALSE;
   BenchUut14.GripButton := FALSE;
   BenchUut14.ReleaseButton := FALSE;
   BenchUut14.DownLimitSwitch := FALSE;
   BenchUut14.UpLimitSwitch := FALSE;
   BenchUut14.LeftLimitSwitch := FALSE;
   BenchUut14.RightLimitSwitch := FALSE;
   BenchUut14.GripLimitSwitch := FALSE;
   BenchUut14.ReleaseLimitSwitch := FALSE;
   TraceIn_ManualMode[170] := BenchUut14.ManualMode;
   TraceIn_SingleStepMode[170] := BenchUut14.SingleStepMode;
   TraceIn_SingleCycleMode[170] := BenchUut14.SingleCycleMode;
   TraceIn_ContinuousMode[170] := BenchUut14.ContinuousMode;
   TraceIn_EmergencyStop[170] := BenchUut14.EmergencyStop;
   TraceIn_Start[170] := BenchUut14.Start;
   TraceIn_DownButton[170] := BenchUut14.DownButton;
   TraceIn_UpButton[170] := BenchUut14.UpButton;
   TraceIn_LeftButton[170] := BenchUut14.LeftButton;
   TraceIn_RightButton[170] := BenchUut14.RightButton;
   TraceIn_GripButton[170] := BenchUut14.GripButton;
   TraceIn_ReleaseButton[170] := BenchUut14.ReleaseButton;
   TraceIn_DownLimitSwitch[170] := BenchUut14.DownLimitSwitch;
   TraceIn_UpLimitSwitch[170] := BenchUut14.UpLimitSwitch;
   TraceIn_LeftLimitSwitch[170] := BenchUut14.LeftLimitSwitch;
   TraceIn_RightLimitSwitch[170] := BenchUut14.RightLimitSwitch;
   TraceIn_GripLimitSwitch[170] := BenchUut14.GripLimitSwitch;
   TraceIn_ReleaseLimitSwitch[170] := BenchUut14.ReleaseLimitSwitch;
   BenchUut14();
   TraceOut_MoveDown[170] := BenchUut14.MoveDown;
   TraceOut_MoveUp[170] := BenchUut14.MoveUp;
   TraceOut_MoveLeft[170] := BenchUut14.MoveLeft;
   TraceOut_MoveRight[170] := BenchUut14.MoveRight;
   TraceOut_ActivateGrip[170] := BenchUut14.ActivateGrip;
   TraceOut_ActivateRelease[170] := BenchUut14.ActivateRelease;
   BenchCalls := BenchCalls + 1;
 171:
   BenchUut14.ManualMode := FALSE;
   BenchUut14.SingleStepMode := TRUE;
   BenchUut14.SingleCycleMode := FALSE;
   BenchUut14.ContinuousMode := FALSE;
   BenchUut14.EmergencyStop := TRUE;
   BenchUut14.Start := FALSE;
   BenchUut14.DownButton := FALSE;
   BenchUut14.UpButton := FALSE;
   BenchUut14.LeftButton := FALSE;
   BenchUut14.RightButton := FALSE;
   BenchUut14.GripButton := FALSE;
   BenchUut14.ReleaseButton := FALSE;
   BenchUut14.DownLimitSwitch := FALSE;
   BenchUut14.UpLimitSwitch := TRUE;
   BenchUut14.LeftLimitSwitch := FALSE;
   BenchUut14.RightLimitSwitch := FALSE;
   BenchUut14.GripLimitSwitch := FALSE;
   BenchUut14.ReleaseLimitSwitch := FALSE;
   TraceIn_ManualMode[171] := BenchUut14.ManualMode;
   TraceIn_SingleStepMode[171] := BenchUut14.SingleStepMode;
   TraceIn_SingleCycleMode[171] := BenchUut14.SingleCycleMode;
   TraceIn_ContinuousMode[171] := BenchUut14.ContinuousMode;
   TraceIn_EmergencyStop[171] := BenchUut14.EmergencyStop;
   TraceIn_Start[171] := BenchUut14.Start;
   TraceIn_DownButton[171] := BenchUut14.DownButton;
   TraceIn_UpButton[171] := BenchUut14.UpButton;
   TraceIn_LeftButton[171] := BenchUut14.LeftButton;
   TraceIn_RightButton[171] := BenchUut14.RightButton;
   TraceIn_GripButton[171] := BenchUut14.GripButton;
   TraceIn_ReleaseButton[171] := BenchUut14.ReleaseButton;
   TraceIn_DownLimitSwitch[171] := BenchUut14.DownLimitSwitch;
   TraceIn_UpLimitSwitch[171] := BenchUut14.UpLimitSwitch;
   TraceIn_LeftLimitSwitch[171] := BenchUut14.LeftLimitSwitch;
   TraceIn_RightLimitSwitch[171] := BenchUut14.RightLimitSwitch;
   TraceIn_GripLimitSwitch[171] := BenchUut14.GripLimitSwitch;
   TraceIn_ReleaseLimitSwitch[171] := BenchUut14.ReleaseLimitSwitch;
   BenchUut14();
   TraceOut_MoveDown[171] := BenchUut14.MoveDown;
   TraceOut_MoveUp[171] := BenchUut14.MoveUp;
   TraceOut_MoveLeft[171] := BenchUut14.MoveLeft;
   TraceOut_MoveRight[171] := BenchUut14.MoveRight;
   TraceOut_ActivateGrip[171] := BenchUut14.ActivateGrip;
   TraceOut_ActivateRelease[171] := BenchUut14.ActivateRelease;
   BenchCalls := BenchCalls + 1;
 172:
   BenchUut14.ManualMode := FALSE;
   BenchUut14.SingleStepMode := TRUE;
   BenchUut14.SingleCycleMode := FALSE;
   BenchUut14.ContinuousMode := FALSE;
   BenchUut14.EmergencyStop := TRUE;
   BenchUut14.Start := TRUE;
   BenchUut14.DownButton := FALSE;
   BenchUut14.UpButton := FALSE;
   BenchUut14.LeftButton := FALSE;
   BenchUut14.RightButton := FALSE;
   BenchUut14.GripButton := FALSE;
   BenchUut14.ReleaseButton := FALSE;
   BenchUut14.DownLimitSwitch := FALSE;
   BenchUut14.UpLimitSwitch := FALSE;
   BenchUut14.LeftLimitSwitch := FALSE;
   BenchUut14.RightLimitSwitch := FALSE;
   BenchUut14.GripLimitSwitch := FALSE;
   BenchUut14.ReleaseLimitSwitch := FALSE;
   TraceIn_ManualMode[172] := BenchUut14.ManualMode;
   TraceIn_SingleStepMode[172] := BenchUut14.SingleStepMode;
   TraceIn_SingleCycleMode[172] := BenchUut14.SingleCycleMode;
   TraceIn_ContinuousMode[172] := BenchUut14.ContinuousMode;
   TraceIn_EmergencyStop[172] := BenchUut14.EmergencyStop;
   TraceIn_Start[172] := BenchUut14.Start;
   TraceIn_DownButton[172] := BenchUut14.DownButton;
   TraceIn_UpButton[172] := BenchUut14.UpButton;
   TraceIn_LeftButton[172] := BenchUut14.LeftButton;
   TraceIn_RightButton[172] := BenchUut14.RightButton;
   TraceIn_GripButton[172] := BenchUut14.GripButton;
   TraceIn_ReleaseButton[172] := BenchUut14.ReleaseButton;
   TraceIn_DownLimitSwitch[172] := BenchUut14.DownLimitSwitch;
   TraceIn_UpLimitSwitch[172] := BenchUut14.UpLimitSwitch;
   TraceIn_LeftLimitSwitch[172] := BenchUut14.LeftLimitSwitch;
   TraceIn_RightLimitSwitch[172] := BenchUut14.RightLimitSwitch;
   TraceIn_GripLimitSwitch[172] := BenchUut14.GripLimitSwitch;
   TraceIn_ReleaseLimitSwitch[172] := BenchUut14.ReleaseLimitSwitch;
   BenchUut14();
   TraceOut_MoveDown[172] := BenchUut14.MoveDown;
   TraceOut_MoveUp[172] := BenchUut14.MoveUp;
   TraceOut_MoveLeft[172] := BenchUut14.MoveLeft;
   TraceOut_MoveRight[172] := BenchUut14.MoveRight;
   TraceOut_ActivateGrip[172] := BenchUut14.ActivateGrip;
   TraceOut_ActivateRelease[172] := BenchUut14.ActivateRelease;
   BenchCalls := BenchCalls + 1;
 173:
   BenchUut14.ManualMode := FALSE;
   BenchUut14.SingleStepMode := TRUE;
   BenchUut14.SingleCycleMode := FALSE;
   BenchUut14.ContinuousMode := FALSE;
   BenchUut14.EmergencyStop := TRUE;
   BenchUut14.Start := FALSE;
   BenchUut14.DownButton := FALSE;
   BenchUut14.UpButton := FALSE;
   BenchUut14.LeftButton := FALSE;
   BenchUut14.RightButton := FALSE;
   BenchUut14.GripButton := FALSE;
   BenchUut14.ReleaseButton := FALSE;
   BenchUut14.DownLimitSwitch := FALSE;
   BenchUut14.UpLimitSwitch := FALSE;
   BenchUut14.LeftLimitSwitch := FALSE;
   BenchUut14.RightLimitSwitch := FALSE;
   BenchUut14.GripLimitSwitch := FALSE;
   BenchUut14.ReleaseLimitSwitch := FALSE;
   TraceIn_ManualMode[173] := BenchUut14.ManualMode;
   TraceIn_SingleStepMode[173] := BenchUut14.SingleStepMode;
   TraceIn_SingleCycleMode[173] := BenchUut14.SingleCycleMode;
   TraceIn_ContinuousMode[173] := BenchUut14.ContinuousMode;
   TraceIn_EmergencyStop[173] := BenchUut14.EmergencyStop;
   TraceIn_Start[173] := BenchUut14.Start;
   TraceIn_DownButton[173] := BenchUut14.DownButton;
   TraceIn_UpButton[173] := BenchUut14.UpButton;
   TraceIn_LeftButton[173] := BenchUut14.LeftButton;
   TraceIn_RightButton[173] := BenchUut14.RightButton;
   TraceIn_GripButton[173] := BenchUut14.GripButton;
   TraceIn_ReleaseButton[173] := BenchUut14.ReleaseButton;
   TraceIn_DownLimitSwitch[173] := BenchUut14.DownLimitSwitch;
   TraceIn_UpLimitSwitch[173] := BenchUut14.UpLimitSwitch;
   TraceIn_LeftLimitSwitch[173] := BenchUut14.LeftLimitSwitch;
   TraceIn_RightLimitSwitch[173] := BenchUut14.RightLimitSwitch;
   TraceIn_GripLimitSwitch[173] := BenchUut14.GripLimitSwitch;
   TraceIn_ReleaseLimitSwitch[173] := BenchUut14.ReleaseLimitSwitch;
   BenchUut14();
   TraceOut_MoveDown[173] := BenchUut14.MoveDown;
   TraceOut_MoveUp[173] := BenchUut14.MoveUp;
   TraceOut_MoveLeft[173] := BenchUut14.MoveLeft;
   TraceOut_MoveRight[173] := BenchUut14.MoveRight;
   TraceOut_ActivateGrip[173] := BenchUut14.ActivateGrip;
   TraceOut_ActivateRelease[173] := BenchUut14.ActivateRelease;
   BenchCalls := BenchCalls + 1;
 174:
   BenchUut14.ManualMode := FALSE;
   BenchUut14.SingleStepMode := TRUE;
   BenchUut14.SingleCycleMode := FALSE;
   BenchUut14.ContinuousMode := FALSE;
   BenchUut14.EmergencyStop := TRUE;
   BenchUut14.Start := FALSE;
   BenchUut14.DownButton := FALSE;
   BenchUut14.UpButton := FALSE;
   BenchUut14.LeftButton := FALSE;
   BenchUut14.RightButton := FALSE;
   BenchUut14.GripButton := FALSE;
   BenchUut14.ReleaseButton := FALSE;
   BenchUut14.DownLimitSwitch := FALSE;
   BenchUut14.UpLimitSwitch := FALSE;
   BenchUut14.LeftLimitSwitch := FALSE;
   BenchUut14.RightLimitSwitch := FALSE;
   BenchUut14.GripLimitSwitch := FALSE;
   BenchUut14.ReleaseLimitSwitch := FALSE;
   TraceIn_ManualMode[174] := BenchUut14.ManualMode;
   TraceIn_SingleStepMode[174] := BenchUut14.SingleStepMode;
   TraceIn_SingleCycleMode[174] := BenchUut14.SingleCycleMode;
   TraceIn_ContinuousMode[174] := BenchUut14.ContinuousMode;
   TraceIn_EmergencyStop[174] := BenchUut14.EmergencyStop;
   TraceIn_Start[174] := BenchUut14.Start;
   TraceIn_DownButton[174] := BenchUut14.DownButton;
   TraceIn_UpButton[174] := BenchUut14.UpButton;
   TraceIn_LeftButton[174] := BenchUut14.LeftButton;
   TraceIn_RightButton[174] := BenchUut14.RightButton;
   TraceIn_GripButton[174] := BenchUut14.GripButton;
   TraceIn_ReleaseButton[174] := BenchUut14.ReleaseButton;
   TraceIn_DownLimitSwitch[174] := BenchUut14.DownLimitSwitch;
   TraceIn_UpLimitSwitch[174] := BenchUut14.UpLimitSwitch;
   TraceIn_LeftLimitSwitch[174] := BenchUut14.LeftLimitSwitch;
   TraceIn_RightLimitSwitch[174] := BenchUut14.RightLimitSwitch;
   TraceIn_GripLimitSwitch[174] := BenchUut14.GripLimitSwitch;
   TraceIn_ReleaseLimitSwitch[174] := BenchUut14.ReleaseLimitSwitch;
   BenchUut14();
   TraceOut_MoveDown[174] := BenchUut14.MoveDown;
   TraceOut_MoveUp[174] := BenchUut14.MoveUp;
   TraceOut_MoveLeft[174] := BenchUut14.MoveLeft;
   TraceOut_MoveRight[174] := BenchUut14.MoveRight;
   TraceOut_ActivateGrip[174] := BenchUut14.ActivateGrip;
   TraceOut_ActivateRelease[174] := BenchUut14.ActivateRelease;
   BenchCalls := BenchCalls + 1;
 175:
   BenchUut14.ManualMode := FALSE;
   BenchUut14.SingleStepMode := TRUE;
   BenchUut14.SingleCycleMode := FALSE;
   BenchUut14.ContinuousMode := FALSE;
   BenchUut14.EmergencyStop := TRUE;
   BenchUut14.Start := FALSE;
   BenchUut14.DownButton := FALSE;
   BenchUut14.UpButton := FALSE;
   BenchUut14.LeftButton := FALSE;
   BenchUut14.RightButton := FALSE;
   BenchUut14.GripButton := FALSE;
   BenchUut14.ReleaseButton := FALSE;
   BenchUut14.DownLimitSwitch := FALSE;
   BenchUut14.UpLimitSwitch := FALSE;
   BenchUut14.LeftLimitSwitch := TRUE;
   BenchUut14.RightLimitSwitch := FALSE;
   BenchUut14.GripLimitSwitch := FALSE;
   BenchUut14.ReleaseLimitSwitch := FALSE;
   TraceIn_ManualMode[175] := BenchUut14.ManualMode;
   TraceIn_SingleStepMode[175] := BenchUut14.SingleStepMode;
   TraceIn_SingleCycleMode[175] := BenchUut14.SingleCycleMode;
   TraceIn_ContinuousMode[175] := BenchUut14.ContinuousMode;
   TraceIn_EmergencyStop[175] := BenchUut14.EmergencyStop;
   TraceIn_Start[175] := BenchUut14.Start;
   TraceIn_DownButton[175] := BenchUut14.DownButton;
   TraceIn_UpButton[175] := BenchUut14.UpButton;
   TraceIn_LeftButton[175] := BenchUut14.LeftButton;
   TraceIn_RightButton[175] := BenchUut14.RightButton;
   TraceIn_GripButton[175] := BenchUut14.GripButton;
   TraceIn_ReleaseButton[175] := BenchUut14.ReleaseButton;
   TraceIn_DownLimitSwitch[175] := BenchUut14.DownLimitSwitch;
   TraceIn_UpLimitSwitch[175] := BenchUut14.UpLimitSwitch;
   TraceIn_LeftLimitSwitch[175] := BenchUut14.LeftLimitSwitch;
   TraceIn_RightLimitSwitch[175] := BenchUut14.RightLimitSwitch;
   TraceIn_GripLimitSwitch[175] := BenchUut14.GripLimitSwitch;
   TraceIn_ReleaseLimitSwitch[175] := BenchUut14.ReleaseLimitSwitch;
   BenchUut14();
   TraceOut_MoveDown[175] := BenchUut14.MoveDown;
   TraceOut_MoveUp[175] := BenchUut14.MoveUp;
   TraceOut_MoveLeft[175] := BenchUut14.MoveLeft;
   TraceOut_MoveRight[175] := BenchUut14.MoveRight;
   TraceOut_ActivateGrip[175] := BenchUut14.ActivateGrip;
   TraceOut_ActivateRelease[175] := BenchUut14.ActivateRelease;
   BenchCalls := BenchCalls + 1;
 176:
   BenchUut15.ManualMode := FALSE;
   BenchUut15.SingleStepMode := FALSE;
   BenchUut15.SingleCycleMode := TRUE;
   BenchUut15.ContinuousMode := FALSE;
   BenchUut15.EmergencyStop := TRUE;
   BenchUut15.Start := FALSE;
   BenchUut15.DownButton := FALSE;
   BenchUut15.UpButton := FALSE;
   BenchUut15.LeftButton := FALSE;
   BenchUut15.RightButton := FALSE;
   BenchUut15.GripButton := FALSE;
   BenchUut15.ReleaseButton := FALSE;
   BenchUut15.DownLimitSwitch := FALSE;
   BenchUut15.UpLimitSwitch := TRUE;
   BenchUut15.LeftLimitSwitch := TRUE;
   BenchUut15.RightLimitSwitch := FALSE;
   BenchUut15.GripLimitSwitch := FALSE;
   BenchUut15.ReleaseLimitSwitch := FALSE;
   TraceIn_ManualMode[176] := BenchUut15.ManualMode;
   TraceIn_SingleStepMode[176] := BenchUut15.SingleStepMode;
   TraceIn_SingleCycleMode[176] := BenchUut15.SingleCycleMode;
   TraceIn_ContinuousMode[176] := BenchUut15.ContinuousMode;
   TraceIn_EmergencyStop[176] := BenchUut15.EmergencyStop;
   TraceIn_Start[176] := BenchUut15.Start;
   TraceIn_DownButton[176] := BenchUut15.DownButton;
   TraceIn_UpButton[176] := BenchUut15.UpButton;
   TraceIn_LeftButton[176] := BenchUut15.LeftButton;
   TraceIn_RightButton[176] := BenchUut15.RightButton;
   TraceIn_GripButton[176] := BenchUut15.GripButton;
   TraceIn_ReleaseButton[176] := BenchUut15.ReleaseButton;
   TraceIn_DownLimitSwitch[176] := BenchUut15.DownLimitSwitch;
   TraceIn_UpLimitSwitch[176] := BenchUut15.UpLimitSwitch;
   TraceIn_LeftLimitSwitch[176] := BenchUut15.LeftLimitSwitch;
   TraceIn_RightLimitSwitch[176] := BenchUut15.RightLimitSwitch;
   TraceIn_GripLimitSwitch[176] := BenchUut15.GripLimitSwitch;
   TraceIn_ReleaseLimitSwitch[176] := BenchUut15.ReleaseLimitSwitch;
   BenchUut15();
   TraceOut_MoveDown[176] := BenchUut15.MoveDown;
   TraceOut_MoveUp[176] := BenchUut15.MoveUp;
   TraceOut_MoveLeft[176] := BenchUut15.MoveLeft;
   TraceOut_MoveRight[176] := BenchUut15.MoveRight;
   TraceOut_ActivateGrip[176] := BenchUut15.ActivateGrip;
   TraceOut_ActivateRelease[176] := BenchUut15.ActivateRelease;
   BenchCalls := BenchCalls + 1;
 177:
   BenchUut15.ManualMode := FALSE;
   BenchUut15.SingleStepMode := FALSE;
   BenchUut15.SingleCycleMode := TRUE;
   BenchUut15.ContinuousMode := FALSE;
   BenchUut15.EmergencyStop := TRUE;
   BenchUut15.Start := TRUE;
   BenchUut15.DownButton := FALSE;
   BenchUut15.UpButton := FALSE;
   BenchUut15.LeftButton := FALSE;
   BenchUut15.RightButton := FALSE;
   BenchUut15.GripButton := FALSE;
   BenchUut15.ReleaseButton := FALSE;
   BenchUut15.DownLimitSwitch := FALSE;
   BenchUut15.UpLimitSwitch := TRUE;
   BenchUut15.LeftLimitSwitch := TRUE;
   BenchUut15.RightLimitSwitch := FALSE;
   BenchUut15.GripLimitSwitch := FALSE;
   BenchUut15.ReleaseLimitSwitch := FALSE;
   TraceIn_ManualMode[177] := BenchUut15.ManualMode;
   TraceIn_SingleStepMode[177] := BenchUut15.SingleStepMode;
   TraceIn_SingleCycleMode[177] := BenchUut15.SingleCycleMode;
   TraceIn_ContinuousMode[177] := BenchUut15.ContinuousMode;
   TraceIn_EmergencyStop[177] := BenchUut15.EmergencyStop;
   TraceIn_Start[177] := BenchUut15.Start;
   TraceIn_DownButton[177] := BenchUut15.DownButton;
   TraceIn_UpButton[177] := BenchUut15.UpButton;
   TraceIn_LeftButton[177] := BenchUut15.LeftButton;
   TraceIn_RightButton[177] := BenchUut15.RightButton;
   TraceIn_GripButton[177] := BenchUut15.GripButton;
   TraceIn_ReleaseButton[177] := BenchUut15.ReleaseButton;
   TraceIn_DownLimitSwitch[177] := BenchUut15.DownLimitSwitch;
   TraceIn_UpLimitSwitch[177] := BenchUut15.UpLimitSwitch;
   TraceIn_LeftLimitSwitch[177] := BenchUut15.LeftLimitSwitch;
   TraceIn_RightLimitSwitch[177] := BenchUut15.RightLimitSwitch;
   TraceIn_GripLimitSwitch[177] := BenchUut15.GripLimitSwitch;
   TraceIn_ReleaseLimitSwitch[177] := BenchUut15.ReleaseLimitSwitch;
   BenchUut15();
   TraceOut_MoveDown[177] := BenchUut15.MoveDown;
   TraceOut_MoveUp[177] := BenchUut15.MoveUp;
   TraceOut_MoveLeft[177] := BenchUut15.MoveLeft;
   TraceOut_MoveRight[177] := BenchUut15.MoveRight;
   TraceOut_ActivateGrip[177] := BenchUut15.ActivateGrip;
   TraceOut_ActivateRelease[177] := BenchUut15.ActivateRelease;
   BenchCalls := BenchCalls + 1;
 178:
   BenchUut15.ManualMode := FALSE;
   BenchUut15.SingleStepMode := FALSE;
   BenchUut15.SingleCycleMode := TRUE;
   BenchUut15.ContinuousMode := FALSE;
   BenchUut15.EmergencyStop := TRUE;
   BenchUut15.Start := FALSE;
   BenchUut15.DownButton := FALSE;
   BenchUut15.UpButton := FALSE;
   BenchUut15.LeftButton := FALSE;
   BenchUut15.RightButton := FALSE;
   BenchUut15.GripButton := FALSE;
   BenchUut15.ReleaseButton := FALSE;
   BenchUut15.DownLimitSwitch := FALSE;
   BenchUut15.UpLimitSwitch := TRUE;
   BenchUut15.LeftLimitSwitch := TRUE;
   BenchUut15.RightLimitSwitch := FALSE;
   BenchUut15.GripLimitSwitch := FALSE;
   BenchUut15.ReleaseLimitSwitch := FALSE;
   TraceIn_ManualMode[178] := BenchUut15.ManualMode;
   TraceIn_SingleStepMode[178] := BenchUut15.SingleStepMode;
   TraceIn_SingleCycleMode[178] := BenchUut15.SingleCycleMode;
   TraceIn_ContinuousMode[178] := BenchUut15.ContinuousMode;
   TraceIn_EmergencyStop[178] := BenchUut15.EmergencyStop;
   TraceIn_Start[178] := BenchUut15.Start;
   TraceIn_DownButton[178] := BenchUut15.DownButton;
   TraceIn_UpButton[178] := BenchUut15.UpButton;
   TraceIn_LeftButton[178] := BenchUut15.LeftButton;
   TraceIn_RightButton[178] := BenchUut15.RightButton;
   TraceIn_GripButton[178] := BenchUut15.GripButton;
   TraceIn_ReleaseButton[178] := BenchUut15.ReleaseButton;
   TraceIn_DownLimitSwitch[178] := BenchUut15.DownLimitSwitch;
   TraceIn_UpLimitSwitch[178] := BenchUut15.UpLimitSwitch;
   TraceIn_LeftLimitSwitch[178] := BenchUut15.LeftLimitSwitch;
   TraceIn_RightLimitSwitch[178] := BenchUut15.RightLimitSwitch;
   TraceIn_GripLimitSwitch[178] := BenchUut15.GripLimitSwitch;
   TraceIn_ReleaseLimitSwitch[178] := BenchUut15.ReleaseLimitSwitch;
   BenchUut15();
   TraceOut_MoveDown[178] := BenchUut15.MoveDown;
   TraceOut_MoveUp[178] := BenchUut15.MoveUp;
   TraceOut_MoveLeft[178] := BenchUut15.MoveLeft;
   TraceOut_MoveRight[178] := BenchUut15.MoveRight;
   TraceOut_ActivateGrip[178] := BenchUut15.ActivateGrip;
   TraceOut_ActivateRelease[178] := BenchUut15.ActivateRelease;
   BenchCalls := BenchCalls + 1;
 179:
   BenchUut15.ManualMode := FALSE;
   BenchUut15.SingleStepMode := FALSE;
   BenchUut15.SingleCycleMode := TRUE;
   BenchUut15.ContinuousMode := FALSE;
   BenchUut15.EmergencyStop := TRUE;
   BenchUut15.Start := FALSE;
   BenchUut15.DownButton := FALSE;
   BenchUut15.UpButton := FALSE;
   BenchUut15.LeftButton := FALSE;
   BenchUut15.RightButton := FALSE;
   BenchUut15.GripButton := FALSE;
   BenchUut15.ReleaseButton := FALSE;
   BenchUut15.DownLimitSwitch := FALSE;
   BenchUut15.UpLimitSwitch := TRUE;
   BenchUut15.LeftLimitSwitch := TRUE;
   BenchUut15.RightLimitSwitch := FALSE;
   BenchUut15.GripLimitSwitch := FALSE;
   BenchUut15.ReleaseLimitSwitch := FALSE;
   TraceIn_ManualMode[179] := BenchUut15.ManualMode;
   TraceIn_SingleStepMode[179] := BenchUut15.SingleStepMode;
   TraceIn_SingleCycleMode[179] := BenchUut15.SingleCycleMode;
   TraceIn_ContinuousMode[179] := BenchUut15.ContinuousMode;
   TraceIn_EmergencyStop[179] := BenchUut15.EmergencyStop;
   TraceIn_Start[179] := BenchUut15.Start;
   TraceIn_DownButton[179] := BenchUut15.DownButton;
   TraceIn_UpButton[179] := BenchUut15.UpButton;
   TraceIn_LeftButton[179] := BenchUut15.LeftButton;
   TraceIn_RightButton[179] := BenchUut15.RightButton;
   TraceIn_GripButton[179] := BenchUut15.GripButton;
   TraceIn_ReleaseButton[179] := BenchUut15.ReleaseButton;
   TraceIn_DownLimitSwitch[179] := BenchUut15.DownLimitSwitch;
   TraceIn_UpLimitSwitch[179] := BenchUut15.UpLimitSwitch;
   TraceIn_LeftLimitSwitch[179] := BenchUut15.LeftLimitSwitch;
   TraceIn_RightLimitSwitch[179] := BenchUut15.RightLimitSwitch;
   TraceIn_GripLimitSwitch[179] := BenchUut15.GripLimitSwitch;
   TraceIn_ReleaseLimitSwitch[179] := BenchUut15.ReleaseLimitSwitch;
   BenchUut15();
   TraceOut_MoveDown[179] := BenchUut15.MoveDown;
   TraceOut_MoveUp[179] := BenchUut15.MoveUp;
   TraceOut_MoveLeft[179] := BenchUut15.MoveLeft;
   TraceOut_MoveRight[179] := BenchUut15.MoveRight;
   TraceOut_ActivateGrip[179] := BenchUut15.ActivateGrip;
   TraceOut_ActivateRelease[179] := BenchUut15.ActivateRelease;
   BenchCalls := BenchCalls + 1;
 180:
   BenchUut15.ManualMode := FALSE;
   BenchUut15.SingleStepMode := FALSE;
   BenchUut15.SingleCycleMode := TRUE;
   BenchUut15.ContinuousMode := FALSE;
   BenchUut15.EmergencyStop := TRUE;
   BenchUut15.Start := FALSE;
   BenchUut15.DownButton := FALSE;
   BenchUut15.UpButton := FALSE;
   BenchUut15.LeftButton := FALSE;
   BenchUut15.RightButton := FALSE;
   BenchUut15.GripButton := FALSE;
   BenchUut15.ReleaseButton := FALSE;
   BenchUut15.DownLimitSwitch := TRUE;
   BenchUut15.UpLimitSwitch := FALSE;
   BenchUut15.LeftLimitSwitch := FALSE;
   BenchUut15.RightLimitSwitch := FALSE;
   BenchUut15.GripLimitSwitch := FALSE;
   BenchUut15.ReleaseLimitSwitch := FALSE;
   TraceIn_ManualMode[180] := BenchUut15.ManualMode;
   TraceIn_SingleStepMode[180] := BenchUut15.SingleStepMode;
   TraceIn_SingleCycleMode[180] := BenchUut15.SingleCycleMode;
   TraceIn_ContinuousMode[180] := BenchUut15.ContinuousMode;
   TraceIn_EmergencyStop[180] := BenchUut15.EmergencyStop;
   TraceIn_Start[180] := BenchUut15.Start;
   TraceIn_DownButton[180] := BenchUut15.DownButton;
   TraceIn_UpButton[180] := BenchUut15.UpButton;
   TraceIn_LeftButton[180] := BenchUut15.LeftButton;
   TraceIn_RightButton[180] := BenchUut15.RightButton;
   TraceIn_GripButton[180] := BenchUut15.GripButton;
   TraceIn_ReleaseButton[180] := BenchUut15.ReleaseButton;
   TraceIn_DownLimitSwitch[180] := BenchUut15.DownLimitSwitch;
   TraceIn_UpLimitSwitch[180] := BenchUut15.UpLimitSwitch;
   TraceIn_LeftLimitSwitch[180] := BenchUut15.LeftLimitSwitch;
   TraceIn_RightLimitSwitch[180] := BenchUut15.RightLimitSwitch;
   TraceIn_GripLimitSwitch[180] := BenchUut15.GripLimitSwitch;
   TraceIn_ReleaseLimitSwitch[180] := BenchUut15.ReleaseLimitSwitch;
   BenchUut15();
   TraceOut_MoveDown[180] := BenchUut15.MoveDown;
   TraceOut_MoveUp[180] := BenchUut15.MoveUp;
   TraceOut_MoveLeft[180] := BenchUut15.MoveLeft;
   TraceOut_MoveRight[180] := BenchUut15.MoveRight;
   TraceOut_ActivateGrip[180] := BenchUut15.ActivateGrip;
   TraceOut_ActivateRelease[180] := BenchUut15.ActivateRelease;
   BenchCalls := BenchCalls + 1;
 181:
   BenchUut15.ManualMode := FALSE;
   BenchUut15.SingleStepMode := FALSE;
   BenchUut15.SingleCycleMode := TRUE;
   BenchUut15.ContinuousMode := FALSE;
   BenchUut15.EmergencyStop := TRUE;
   BenchUut15.Start := FALSE;
   BenchUut15.DownButton := FALSE;
   BenchUut15.UpButton := FALSE;
   BenchUut15.LeftButton := FALSE;
   BenchUut15.RightButton := FALSE;
   BenchUut15.GripButton := FALSE;
   BenchUut15.ReleaseButton := FALSE;
   BenchUut15.DownLimitSwitch := FALSE;
   BenchUut15.UpLimitSwitch := FALSE;
   BenchUut15.LeftLimitSwitch := FALSE;
   BenchUut15.RightLimitSwitch := FALSE;
   BenchUut15.GripLimitSwitch := FALSE;
   BenchUut15.ReleaseLimitSwitch := FALSE;
   TraceIn_ManualMode[181] := BenchUut15.ManualMode;
   TraceIn_SingleStepMode[181] := BenchUut15.SingleStepMode;
   TraceIn_SingleCycleMode[181] := BenchUut15.SingleCycleMode;
   TraceIn_ContinuousMode[181] := BenchUut15.ContinuousMode;
   TraceIn_EmergencyStop[181] := BenchUut15.EmergencyStop;
   TraceIn_Start[181] := BenchUut15.Start;
   TraceIn_DownButton[181] := BenchUut15.DownButton;
   TraceIn_UpButton[181] := BenchUut15.UpButton;
   TraceIn_LeftButton[181] := BenchUut15.LeftButton;
   TraceIn_RightButton[181] := BenchUut15.RightButton;
   TraceIn_GripButton[181] := BenchUut15.GripButton;
   TraceIn_ReleaseButton[181] := BenchUut15.ReleaseButton;
   TraceIn_DownLimitSwitch[181] := BenchUut15.DownLimitSwitch;
   TraceIn_UpLimitSwitch[181] := BenchUut15.UpLimitSwitch;
   TraceIn_LeftLimitSwitch[181] := BenchUut15.LeftLimitSwitch;
   TraceIn_RightLimitSwitch[181] := BenchUut15.RightLimitSwitch;
   TraceIn_GripLimitSwitch[181] := BenchUut15.GripLimitSwitch;
   TraceIn_ReleaseLimitSwitch[181] := BenchUut15.ReleaseLimitSwitch;
   BenchUut15();
   TraceOut_MoveDown[181] := BenchUut15.MoveDown;
   TraceOut_MoveUp[181] := BenchUut15.MoveUp;
   TraceOut_MoveLeft[181] := BenchUut15.MoveLeft;
   TraceOut_MoveRight[181] := BenchUut15.MoveRight;
   TraceOut_ActivateGrip[181] := BenchUut15.ActivateGrip;
   TraceOut_ActivateRelease[181] := BenchUut15.ActivateRelease;
   BenchCalls := BenchCalls + 1;
 182:
   BenchUut15.ManualMode := FALSE;
   BenchUut15.SingleStepMode := FALSE;
   BenchUut15.SingleCycleMode := TRUE;
   BenchUut15.ContinuousMode := FALSE;
   BenchUut15.EmergencyStop := TRUE;
   BenchUut15.Start := FALSE;
   BenchUut15.DownButton := FALSE;
   BenchUut15.UpButton := FALSE;
   BenchUut15.LeftButton := FALSE;
   BenchUut15.RightButton := FALSE;
   BenchUut15.GripButton := FALSE;
   BenchUut15.ReleaseButton := FALSE;
   BenchUut15.DownLimitSwitch := FALSE;
   BenchUut15.UpLimitSwitch := FALSE;
   BenchUut15.LeftLimitSwitch := FALSE;
   BenchUut15.RightLimitSwitch := FALSE;
   BenchUut15.GripLimitSwitch := FALSE;
   BenchUut15.ReleaseLimitSwitch := FALSE;
   TraceIn_ManualMode[182] := BenchUut15.ManualMode;
   TraceIn_SingleStepMode[182] := BenchUut15.SingleStepMode;
   TraceIn_SingleCycleMode[182] := BenchUut15.SingleCycleMode;
   TraceIn_ContinuousMode[182] := BenchUut15.ContinuousMode;
   TraceIn_EmergencyStop[182] := BenchUut15.EmergencyStop;
   TraceIn_Start[182] := BenchUut15.Start;
   TraceIn_DownButton[182] := BenchUut15.DownButton;
   TraceIn_UpButton[182] := BenchUut15.UpButton;
   TraceIn_LeftButton[182] := BenchUut15.LeftButton;
   TraceIn_RightButton[182] := BenchUut15.RightButton;
   TraceIn_GripButton[182] := BenchUut15.GripButton;
   TraceIn_ReleaseButton[182] := BenchUut15.ReleaseButton;
   TraceIn_DownLimitSwitch[182] := BenchUut15.DownLimitSwitch;
   TraceIn_UpLimitSwitch[182] := BenchUut15.UpLimitSwitch;
   TraceIn_LeftLimitSwitch[182] := BenchUut15.LeftLimitSwitch;
   TraceIn_RightLimitSwitch[182] := BenchUut15.RightLimitSwitch;
   TraceIn_GripLimitSwitch[182] := BenchUut15.GripLimitSwitch;
   TraceIn_ReleaseLimitSwitch[182] := BenchUut15.ReleaseLimitSwitch;
   BenchUut15();
   TraceOut_MoveDown[182] := BenchUut15.MoveDown;
   TraceOut_MoveUp[182] := BenchUut15.MoveUp;
   TraceOut_MoveLeft[182] := BenchUut15.MoveLeft;
   TraceOut_MoveRight[182] := BenchUut15.MoveRight;
   TraceOut_ActivateGrip[182] := BenchUut15.ActivateGrip;
   TraceOut_ActivateRelease[182] := BenchUut15.ActivateRelease;
   BenchCalls := BenchCalls + 1;
 183:
   BenchUut15.ManualMode := FALSE;
   BenchUut15.SingleStepMode := FALSE;
   BenchUut15.SingleCycleMode := TRUE;
   BenchUut15.ContinuousMode := FALSE;
   BenchUut15.EmergencyStop := TRUE;
   BenchUut15.Start := FALSE;
   BenchUut15.DownButton := FALSE;
   BenchUut15.UpButton := FALSE;
   BenchUut15.LeftButton := FALSE;
   BenchUut15.RightButton := FALSE;
   BenchUut15.GripButton := FALSE;
   BenchUut15.ReleaseButton := FALSE;
   BenchUut15.DownLimitSwitch := FALSE;
   BenchUut15.UpLimitSwitch := FALSE;
   BenchUut15.LeftLimitSwitch := FALSE;
   BenchUut15.RightLimitSwitch := FALSE;
   BenchUut15.GripLimitSwitch := FALSE;
   BenchUut15.ReleaseLimitSwitch := FALSE;
   TraceIn_ManualMode[183] := BenchUut15.ManualMode;
   TraceIn_SingleStepMode[183] := BenchUut15.SingleStepMode;
   TraceIn_SingleCycleMode[183] := BenchUut15.SingleCycleMode;
   TraceIn_ContinuousMode[183] := BenchUut15.ContinuousMode;
   TraceIn_EmergencyStop[183] := BenchUut15.EmergencyStop;
   TraceIn_Start[183] := BenchUut15.Start;
   TraceIn_DownButton[183] := BenchUut15.DownButton;
   TraceIn_UpButton[183] := BenchUut15.UpButton;
   TraceIn_LeftButton[183] := BenchUut15.LeftButton;
   TraceIn_RightButton[183] := BenchUut15.RightButton;
   TraceIn_GripButton[183] := BenchUut15.GripButton;
   TraceIn_ReleaseButton[183] := BenchUut15.ReleaseButton;
   TraceIn_DownLimitSwitch[183] := BenchUut15.DownLimitSwitch;
   TraceIn_UpLimitSwitch[183] := BenchUut15.UpLimitSwitch;
   TraceIn_LeftLimitSwitch[183] := BenchUut15.LeftLimitSwitch;
   TraceIn_RightLimitSwitch[183] := BenchUut15.RightLimitSwitch;
   TraceIn_GripLimitSwitch[183] := BenchUut15.GripLimitSwitch;
   TraceIn_ReleaseLimitSwitch[183] := BenchUut15.ReleaseLimitSwitch;
   BenchUut15();
   TraceOut_MoveDown[183] := BenchUut15.MoveDown;
   TraceOut_MoveUp[183] := BenchUut15.MoveUp;
   TraceOut_MoveLeft[183] := BenchUut15.MoveLeft;
   TraceOut_MoveRight[183] := BenchUut15.MoveRight;
   TraceOut_ActivateGrip[183] := BenchUut15.ActivateGrip;
   TraceOut_ActivateRelease[183] := BenchUut15.ActivateRelease;
   BenchCalls := BenchCalls + 1;
 184:
   BenchUut15.ManualMode := FALSE;
   BenchUut15.SingleStepMode := FALSE;
   BenchUut15.SingleCycleMode := TRUE;
   BenchUut15.ContinuousMode := FALSE;
   BenchUut15.EmergencyStop := TRUE;
   BenchUut15.Start := FALSE;
   BenchUut15.DownButton := FALSE;
   BenchUut15.UpButton := FALSE;
   BenchUut15.LeftButton := FALSE;
   BenchUut15.RightButton := FALSE;
   BenchUut15.GripButton := FALSE;
   BenchUut15.ReleaseButton := FALSE;
   BenchUut15.DownLimitSwitch := FALSE;
   BenchUut15.UpLimitSwitch := FALSE;
   BenchUut15.LeftLimitSwitch := FALSE;
   BenchUut15.RightLimitSwitch := FALSE;
   BenchUut15.GripLimitSwitch := TRUE;
   BenchUut15.ReleaseLimitSwitch := FALSE;
   TraceIn_ManualMode[184] := BenchUut15.ManualMode;
   TraceIn_SingleStepMode[184] := BenchUut15.SingleStepMode;
   TraceIn_SingleCycleMode[184] := BenchUut15.SingleCycleMode;
   TraceIn_ContinuousMode[184] := BenchUut15.ContinuousMode;
   TraceIn_EmergencyStop[184] := BenchUut15.EmergencyStop;
   TraceIn_Start[184] := BenchUut15.Start;
   TraceIn_DownButton[184] := BenchUut15.DownButton;
   TraceIn_UpButton[184] := BenchUut15.UpButton;
   TraceIn_LeftButton[184] := BenchUut15.LeftButton;
   TraceIn_RightButton[184] := BenchUut15.RightButton;
   TraceIn_GripButton[184] := BenchUut15.GripButton;
   TraceIn_ReleaseButton[184] := BenchUut15.ReleaseButton;
   TraceIn_DownLimitSwitch[184] := BenchUut15.DownLimitSwitch;
   TraceIn_UpLimitSwitch[184] := BenchUut15.UpLimitSwitch;
   TraceIn_LeftLimitSwitch[184] := BenchUut15.LeftLimitSwitch;
   TraceIn_RightLimitSwitch[184] := BenchUut15.RightLimitSwitch;
   TraceIn_GripLimitSwitch[184] := BenchUut15.GripLimitSwitch;
   TraceIn_ReleaseLimitSwitch[184] := BenchUut15.ReleaseLimitSwitch;
   BenchUut15();
   TraceOut_MoveDown[184] := BenchUut15.MoveDown;
   TraceOut_MoveUp[184] := BenchUut15.MoveUp;
   TraceOut_MoveLeft[184] := BenchUut15.MoveLeft;
   TraceOut_MoveRight[184] := BenchUut15.MoveRight;
   TraceOut_ActivateGrip[184] := BenchUut15.ActivateGrip;
   TraceOut_ActivateRelease[184] := BenchUut15.ActivateRelease;
   BenchCalls := BenchCalls + 1;
 185:
   BenchUut15.ManualMode := FALSE;
   BenchUut15.SingleStepMode := FALSE;
   BenchUut15.SingleCycleMode := TRUE;
   BenchUut15.ContinuousMode := FALSE;
   BenchUut15.EmergencyStop := TRUE;
   BenchUut15.Start := FALSE;
   BenchUut15.DownButton := FALSE;
   BenchUut15.UpButton := FALSE;
   BenchUut15.LeftButton := FALSE;
   BenchUut15.RightButton := FALSE;
   BenchUut15.GripButton := FALSE;
   BenchUut15.ReleaseButton := FALSE;
   BenchUut15.DownLimitSwitch := FALSE;
   BenchUut15.UpLimitSwitch := FALSE;
   BenchUut15.LeftLimitSwitch := FALSE;
   BenchUut15.RightLimitSwitch := FALSE;
   BenchUut15.GripLimitSwitch := FALSE;
   BenchUut15.ReleaseLimitSwitch := FALSE;
   TraceIn_ManualMode[185] := BenchUut15.ManualMode;
   TraceIn_SingleStepMode[185] := BenchUut15.SingleStepMode;
   TraceIn_SingleCycleMode[185] := BenchUut15.SingleCycleMode;
   TraceIn_ContinuousMode[185] := BenchUut15.ContinuousMode;
   TraceIn_EmergencyStop[185] := BenchUut15.EmergencyStop;
   TraceIn_Start[185] := BenchUut15.Start;
   TraceIn_DownButton[185] := BenchUut15.DownButton;
   TraceIn_UpButton[185] := BenchUut15.UpButton;
   TraceIn_LeftButton[185] := BenchUut15.LeftButton;
   TraceIn_RightButton[185] := BenchUut15.RightButton;
   TraceIn_GripButton[185] := BenchUut15.GripButton;
   TraceIn_ReleaseButton[185] := BenchUut15.ReleaseButton;
   TraceIn_DownLimitSwitch[185] := BenchUut15.DownLimitSwitch;
   TraceIn_UpLimitSwitch[185] := BenchUut15.UpLimitSwitch;
   TraceIn_LeftLimitSwitch[185] := BenchUut15.LeftLimitSwitch;
   TraceIn_RightLimitSwitch[185] := BenchUut15.RightLimitSwitch;
   TraceIn_GripLimitSwitch[185] := BenchUut15.GripLimitSwitch;
   TraceIn_ReleaseLimitSwitch[185] := BenchUut15.ReleaseLimitSwitch;
   BenchUut15();
   TraceOut_MoveDown[185] := BenchUut15.MoveDown;
   TraceOut_MoveUp[185] := BenchUut15.MoveUp;
   TraceOut_MoveLeft[185] := BenchUut15.MoveLeft;
   TraceOut_MoveRight[185] := BenchUut15.MoveRight;
   TraceOut_ActivateGrip[185] := BenchUut15.ActivateGrip;
   TraceOut_ActivateRelease[185] := BenchUut15.ActivateRelease;
   BenchCalls := BenchCalls + 1;
 186:
   BenchUut15.ManualMode := FALSE;
   BenchUut15.SingleStepMode := FALSE;
   BenchUut15.SingleCycleMode := TRUE;
   BenchUut15.ContinuousMode := FALSE;
   BenchUut15.EmergencyStop := TRUE;
   BenchUut15.Start := FALSE;
   BenchUut15.DownButton := FALSE;
   BenchUut15.UpButton := FALSE;
   BenchUut15.LeftButton := FALSE;
   BenchUut15.RightButton := FALSE;
   BenchUut15.GripButton := FALSE;
   BenchUut15.ReleaseButton := FALSE;
   BenchUut15.DownLimitSwitch := FALSE;
   BenchUut15.UpLimitSwitch := FALSE;
   BenchUut15.LeftLimitSwitch := FALSE;
   BenchUut15.RightLimitSwitch := FALSE;
   BenchUut15.GripLimitSwitch := FALSE;
   BenchUut15.ReleaseLimitSwitch := FALSE;
   TraceIn_ManualMode[186] := BenchUut15.ManualMode;
   TraceIn_SingleStepMode[186] := BenchUut15.SingleStepMode;
   TraceIn_SingleCycleMode[186] := BenchUut15.SingleCycleMode;
   TraceIn_ContinuousMode[186] := BenchUut15.ContinuousMode;
   TraceIn_EmergencyStop[186] := BenchUut15.EmergencyStop;
   TraceIn_Start[186] := BenchUut15.Start;
   TraceIn_DownButton[186] := BenchUut15.DownButton;
   TraceIn_UpButton[186] := BenchUut15.UpButton;
   TraceIn_LeftButton[186] := BenchUut15.LeftButton;
   TraceIn_RightButton[186] := BenchUut15.RightButton;
   TraceIn_GripButton[186] := BenchUut15.GripButton;
   TraceIn_ReleaseButton[186] := BenchUut15.ReleaseButton;
   TraceIn_DownLimitSwitch[186] := BenchUut15.DownLimitSwitch;
   TraceIn_UpLimitSwitch[186] := BenchUut15.UpLimitSwitch;
   TraceIn_LeftLimitSwitch[186] := BenchUut15.LeftLimitSwitch;
   TraceIn_RightLimitSwitch[186] := BenchUut15.RightLimitSwitch;
   TraceIn_GripLimitSwitch[186] := BenchUut15.GripLimitSwitch;
   TraceIn_ReleaseLimitSwitch[186] := BenchUut15.ReleaseLimitSwitch;
   BenchUut15();
   TraceOut_MoveDown[186] := BenchUut15.MoveDown;
   TraceOut_MoveUp[186] := BenchUut15.MoveUp;
   TraceOut_MoveLeft[186] := BenchUut15.MoveLeft;
   TraceOut_MoveRight[186] := BenchUut15.MoveRight;
   TraceOut_ActivateGrip[186] := BenchUut15.ActivateGrip;
   TraceOut_ActivateRelease[186] := BenchUut15.ActivateRelease;
   BenchCalls := BenchCalls + 1;
 187:
   BenchUut15.ManualMode := FALSE;
   BenchUut15.SingleStepMode := FALSE;
   BenchUut15.SingleCycleMode := TRUE;
   BenchUut15.ContinuousMode := FALSE;
   BenchUut15.EmergencyStop := TRUE;
   BenchUut15.Start := FALSE;
   BenchUut15.DownButton := FALSE;
   BenchUut15.UpButton := FALSE;
   BenchUut15.LeftButton := FALSE;
   BenchUut15.RightButton := FALSE;
   BenchUut15.GripButton := FALSE;
   BenchUut15.ReleaseButton := FALSE;
   BenchUut15.DownLimitSwitch := FALSE;
   BenchUut15.UpLimitSwitch := FALSE;
   BenchUut15.LeftLimitSwitch := FALSE;
   BenchUut15.RightLimitSwitch := FALSE;
   BenchUut15.GripLimitSwitch := FALSE;
   BenchUut15.ReleaseLimitSwitch := FALSE;
   TraceIn_ManualMode[187] := BenchUut15.ManualMode;
   TraceIn_SingleStepMode[187] := BenchUut15.SingleStepMode;
   TraceIn_SingleCycleMode[187] := BenchUut15.SingleCycleMode;
   TraceIn_ContinuousMode[187] := BenchUut15.ContinuousMode;
   TraceIn_EmergencyStop[187] := BenchUut15.EmergencyStop;
   TraceIn_Start[187] := BenchUut15.Start;
   TraceIn_DownButton[187] := BenchUut15.DownButton;
   TraceIn_UpButton[187] := BenchUut15.UpButton;
   TraceIn_LeftButton[187] := BenchUut15.LeftButton;
   TraceIn_RightButton[187] := BenchUut15.RightButton;
   TraceIn_GripButton[187] := BenchUut15.GripButton;
   TraceIn_ReleaseButton[187] := BenchUut15.ReleaseButton;
   TraceIn_DownLimitSwitch[187] := BenchUut15.DownLimitSwitch;
   TraceIn_UpLimitSwitch[187] := BenchUut15.UpLimitSwitch;
   TraceIn_LeftLimitSwitch[187] := BenchUut15.LeftLimitSwitch;
   TraceIn_RightLimitSwitch[187] := BenchUut15.RightLimitSwitch;
   TraceIn_GripLimitSwitch[187] := BenchUut15.GripLimitSwitch;
   TraceIn_ReleaseLimitSwitch[187] := BenchUut15.ReleaseLimitSwitch;
   BenchUut15();
   TraceOut_MoveDown[187] := BenchUut15.MoveDown;
   TraceOut_MoveUp[187] := BenchUut15.MoveUp;
   TraceOut_MoveLeft[187] := BenchUut15.MoveLeft;
   TraceOut_MoveRight[187] := BenchUut15.MoveRight;
   TraceOut_ActivateGrip[187] := BenchUut15.ActivateGrip;
   TraceOut_ActivateRelease[187] := BenchUut15.ActivateRelease;
   BenchCalls := BenchCalls + 1;
 188:
   BenchUut15.ManualMode := FALSE;
   BenchUut15.SingleStepMode := FALSE;
   BenchUut15.SingleCycleMode := TRUE;
   BenchUut15.ContinuousMode := FALSE;
   BenchUut15.EmergencyStop := TRUE;
   BenchUut15.Start := FALSE;
   BenchUut15.DownButton := FALSE;
   BenchUut15.UpButton := FALSE;
   BenchUut15.LeftButton := FALSE;
   BenchUut15.RightButton := FALSE;
   BenchUut15.GripButton := FALSE;
   BenchUut15.ReleaseButton := FALSE;
   BenchUut15.DownLimitSwitch := FALSE;
   BenchUut15.UpLimitSwitch := TRUE;
   BenchUut15.LeftLimitSwitch := FALSE;
   BenchUut15.RightLimitSwitch := FALSE;
   BenchUut15.GripLimitSwitch := FALSE;
   BenchUut15.ReleaseLimitSwitch := FALSE;
   TraceIn_ManualMode[188] := BenchUut15.ManualMode;
   TraceIn_SingleStepMode[188] := BenchUut15.SingleStepMode;
   TraceIn_SingleCycleMode[188] := BenchUut15.SingleCycleMode;
   TraceIn_ContinuousMode[188] := BenchUut15.ContinuousMode;
   TraceIn_EmergencyStop[188] := BenchUut15.EmergencyStop;
   TraceIn_Start[188] := BenchUut15.Start;
   TraceIn_DownButton[188] := BenchUut15.DownButton;
   TraceIn_UpButton[188] := BenchUut15.UpButton;
   TraceIn_LeftButton[188] := BenchUut15.LeftButton;
   TraceIn_RightButton[188] := BenchUut15.RightButton;
   TraceIn_GripButton[188] := BenchUut15.GripButton;
   TraceIn_ReleaseButton[188] := BenchUut15.ReleaseButton;
   TraceIn_DownLimitSwitch[188] := BenchUut15.DownLimitSwitch;
   TraceIn_UpLimitSwitch[188] := BenchUut15.UpLimitSwitch;
   TraceIn_LeftLimitSwitch[188] := BenchUut15.LeftLimitSwitch;
   TraceIn_RightLimitSwitch[188] := BenchUut15.RightLimitSwitch;
   TraceIn_GripLimitSwitch[188] := BenchUut15.GripLimitSwitch;
   TraceIn_ReleaseLimitSwitch[188] := BenchUut15.ReleaseLimitSwitch;
   BenchUut15();
   TraceOut_MoveDown[188] := BenchUut15.MoveDown;
   TraceOut_MoveUp[188] := BenchUut15.MoveUp;
   TraceOut_MoveLeft[188] := BenchUut15.MoveLeft;
   TraceOut_MoveRight[188] := BenchUut15.MoveRight;
   TraceOut_ActivateGrip[188] := BenchUut15.ActivateGrip;
   TraceOut_ActivateRelease[188] := BenchUut15.ActivateRelease;
   BenchCalls := BenchCalls + 1;
 189:
   BenchUut15.ManualMode := FALSE;
   BenchUut15.SingleStepMode := FALSE;
   BenchUut15.SingleCycleMode := TRUE;
   BenchUut15.ContinuousMode := FALSE;
   BenchUut15.EmergencyStop := TRUE;
   BenchUut15.Start := FALSE;
   BenchUut15.DownButton := FALSE;
   BenchUut15.UpButton := FALSE;
   BenchUut15.LeftButton := FALSE;
   BenchUut15.RightButton := FALSE;
   BenchUut15.GripButton := FALSE;
   BenchUut15.ReleaseButton := FALSE;
   BenchUut15.DownLimitSwitch := FALSE;
   BenchUut15.UpLimitSwitch := FALSE;
   BenchUut15.LeftLimitSwitch := FALSE;
   BenchUut15.RightLimitSwitch := FALSE;
   BenchUut15.GripLimitSwitch := FALSE;
   BenchUut15.ReleaseLimitSwitch := FALSE;
   TraceIn_ManualMode[189] := BenchUut15.ManualMode;
   TraceIn_SingleStepMode[189] := BenchUut15.SingleStepMode;
   TraceIn_SingleCycleMode[189] := BenchUut15.SingleCycleMode;
   TraceIn_ContinuousMode[189] := BenchUut15.ContinuousMode;
   TraceIn_EmergencyStop[189] := BenchUut15.EmergencyStop;
   TraceIn_Start[189] := BenchUut15.Start;
   TraceIn_DownButton[189] := BenchUut15.DownButton;
   TraceIn_UpButton[189] := BenchUut15.UpButton;
   TraceIn_LeftButton[189] := BenchUut15.LeftButton;
   TraceIn_RightButton[189] := BenchUut15.RightButton;
   TraceIn_GripButton[189] := BenchUut15.GripButton;
   TraceIn_ReleaseButton[189] := BenchUut15.ReleaseButton;
   TraceIn_DownLimitSwitch[189] := BenchUut15.DownLimitSwitch;
   TraceIn_UpLimitSwitch[189] := BenchUut15.UpLimitSwitch;
   TraceIn_LeftLimitSwitch[189] := BenchUut15.LeftLimitSwitch;
   TraceIn_RightLimitSwitch[189] := BenchUut15.RightLimitSwitch;
   TraceIn_GripLimitSwitch[189] := BenchUut15.GripLimitSwitch;
   TraceIn_ReleaseLimitSwitch[189] := BenchUut15.ReleaseLimitSwitch;
   BenchUut15();
   TraceOut_MoveDown[189] := BenchUut15.MoveDown;
   TraceOut_MoveUp[189] := BenchUut15.MoveUp;
   TraceOut_MoveLeft[189] := BenchUut15.MoveLeft;
   TraceOut_MoveRight[189] := BenchUut15.MoveRight;
   TraceOut_ActivateGrip[189] := BenchUut15.ActivateGrip;
   TraceOut_ActivateRelease[189] := BenchUut15.ActivateRelease;
   BenchCalls := BenchCalls + 1;
 190:
   BenchUut15.ManualMode := FALSE;
   BenchUut15.SingleStepMode := FALSE;
   BenchUut15.SingleCycleMode := TRUE;
   BenchUut15.ContinuousMode := FALSE;
   BenchUut15.EmergencyStop := TRUE;
   BenchUut15.Start := FALSE;
   BenchUut15.DownButton := FALSE;
   BenchUut15.UpButton := FALSE;
   BenchUut15.LeftButton := FALSE;
   BenchUut15.RightButton := FALSE;
   BenchUut15.GripButton := FALSE;
   BenchUut15.ReleaseButton := FALSE;
   BenchUut15.DownLimitSwitch := FALSE;
   BenchUut15.UpLimitSwitch := FALSE;
   BenchUut15.LeftLimitSwitch := FALSE;
   BenchUut15.RightLimitSwitch := FALSE;
   BenchUut15.GripLimitSwitch := FALSE;
   BenchUut15.ReleaseLimitSwitch := FALSE;
   TraceIn_ManualMode[190] := BenchUut15.ManualMode;
   TraceIn_SingleStepMode[190] := BenchUut15.SingleStepMode;
   TraceIn_SingleCycleMode[190] := BenchUut15.SingleCycleMode;
   TraceIn_ContinuousMode[190] := BenchUut15.ContinuousMode;
   TraceIn_EmergencyStop[190] := BenchUut15.EmergencyStop;
   TraceIn_Start[190] := BenchUut15.Start;
   TraceIn_DownButton[190] := BenchUut15.DownButton;
   TraceIn_UpButton[190] := BenchUut15.UpButton;
   TraceIn_LeftButton[190] := BenchUut15.LeftButton;
   TraceIn_RightButton[190] := BenchUut15.RightButton;
   TraceIn_GripButton[190] := BenchUut15.GripButton;
   TraceIn_ReleaseButton[190] := BenchUut15.ReleaseButton;
   TraceIn_DownLimitSwitch[190] := BenchUut15.DownLimitSwitch;
   TraceIn_UpLimitSwitch[190] := BenchUut15.UpLimitSwitch;
   TraceIn_LeftLimitSwitch[190] := BenchUut15.LeftLimitSwitch;
   TraceIn_RightLimitSwitch[190] := BenchUut15.RightLimitSwitch;
   TraceIn_GripLimitSwitch[190] := BenchUut15.GripLimitSwitch;
   TraceIn_ReleaseLimitSwitch[190] := BenchUut15.ReleaseLimitSwitch;
   BenchUut15();
   TraceOut_MoveDown[190] := BenchUut15.MoveDown;
   TraceOut_MoveUp[190] := BenchUut15.MoveUp;
   TraceOut_MoveLeft[190] := BenchUut15.MoveLeft;
   TraceOut_MoveRight[190] := BenchUut15.MoveRight;
   TraceOut_ActivateGrip[190] := BenchUut15.ActivateGrip;
   TraceOut_ActivateRelease[190] := BenchUut15.ActivateRelease;
   BenchCalls := BenchCalls + 1;
 191:
   BenchUut15.ManualMode := FALSE;
   BenchUut15.SingleStepMode := FALSE;
   BenchUut15.SingleCycleMode := TRUE;
   BenchUut15.ContinuousMode := FALSE;
   BenchUut15.EmergencyStop := TRUE;
   BenchUut15.Start := FALSE;
   BenchUut15.DownButton := FALSE;
   BenchUut15.UpButton := FALSE;
   BenchUut15.LeftButton := FALSE;
   BenchUut15.RightButton := FALSE;
   BenchUut15.GripButton := FALSE;
   BenchUut15.ReleaseButton := FALSE;
   BenchUut15.DownLimitSwitch := FALSE;
   BenchUut15.UpLimitSwitch := FALSE;
   BenchUut15.LeftLimitSwitch := FALSE;
   BenchUut15.RightLimitSwitch := FALSE;
   BenchUut15.GripLimitSwitch := FALSE;
   BenchUut15.ReleaseLimitSwitch := FALSE;
   TraceIn_ManualMode[191] := BenchUut15.ManualMode;
   TraceIn_SingleStepMode[191] := BenchUut15.SingleStepMode;
   TraceIn_SingleCycleMode[191] := BenchUut15.SingleCycleMode;
   TraceIn_ContinuousMode[191] := BenchUut15.ContinuousMode;
   TraceIn_EmergencyStop[191] := BenchUut15.EmergencyStop;
   TraceIn_Start[191] := BenchUut15.Start;
   TraceIn_DownButton[191] := BenchUut15.DownButton;
   TraceIn_UpButton[191] := BenchUut15.UpButton;
   TraceIn_LeftButton[191] := BenchUut15.LeftButton;
   TraceIn_RightButton[191] := BenchUut15.RightButton;
   TraceIn_GripButton[191] := BenchUut15.GripButton;
   TraceIn_ReleaseButton[191] := BenchUut15.ReleaseButton;
   TraceIn_DownLimitSwitch[191] := BenchUut15.DownLimitSwitch;
   TraceIn_UpLimitSwitch[191] := BenchUut15.UpLimitSwitch;
   TraceIn_LeftLimitSwitch[191] := BenchUut15.LeftLimitSwitch;
   TraceIn_RightLimitSwitch[191] := BenchUut15.RightLimitSwitch;
   TraceIn_GripLimitSwitch[191] := BenchUut15.GripLimitSwitch;
   TraceIn_ReleaseLimitSwitch[191] := BenchUut15.ReleaseLimitSwitch;
   BenchUut15();
   TraceOut_MoveDown[191] := BenchUut15.MoveDown;
   TraceOut_MoveUp[191] := BenchUut15.MoveUp;
   TraceOut_MoveLeft[191] := BenchUut15.MoveLeft;
   TraceOut_MoveRight[191] := BenchUut15.MoveRight;
   TraceOut_ActivateGrip[191] := BenchUut15.ActivateGrip;
   TraceOut_ActivateRelease[191] := BenchUut15.ActivateRelease;
   BenchCalls := BenchCalls + 1;
 192:
   BenchUut15.ManualMode := FALSE;
   BenchUut15.SingleStepMode := FALSE;
   BenchUut15.SingleCycleMode := TRUE;
   BenchUut15.ContinuousMode := FALSE;
   BenchUut15.EmergencyStop := TRUE;
   BenchUut15.Start := FALSE;
   BenchUut15.DownButton := FALSE;
   BenchUut15.UpButton := FALSE;
   BenchUut15.LeftButton := FALSE;
   BenchUut15.RightButton := FALSE;
   BenchUut15.GripButton := FALSE;
   BenchUut15.ReleaseButton := FALSE;
   BenchUut15.DownLimitSwitch := FALSE;
   BenchUut15.UpLimitSwitch := FALSE;
   BenchUut15.LeftLimitSwitch := FALSE;
   BenchUut15.RightLimitSwitch := TRUE;
   BenchUut15.GripLimitSwitch := FALSE;
   BenchUut15.ReleaseLimitSwitch := FALSE;
   TraceIn_ManualMode[192] := BenchUut15.ManualMode;
   TraceIn_SingleStepMode[192] := BenchUut15.SingleStepMode;
   TraceIn_SingleCycleMode[192] := BenchUut15.SingleCycleMode;
   TraceIn_ContinuousMode[192] := BenchUut15.ContinuousMode;
   TraceIn_EmergencyStop[192] := BenchUut15.EmergencyStop;
   TraceIn_Start[192] := BenchUut15.Start;
   TraceIn_DownButton[192] := BenchUut15.DownButton;
   TraceIn_UpButton[192] := BenchUut15.UpButton;
   TraceIn_LeftButton[192] := BenchUut15.LeftButton;
   TraceIn_RightButton[192] := BenchUut15.RightButton;
   TraceIn_GripButton[192] := BenchUut15.GripButton;
   TraceIn_ReleaseButton[192] := BenchUut15.ReleaseButton;
   TraceIn_DownLimitSwitch[192] := BenchUut15.DownLimitSwitch;
   TraceIn_UpLimitSwitch[192] := BenchUut15.UpLimitSwitch;
   TraceIn_LeftLimitSwitch[192] := BenchUut15.LeftLimitSwitch;
   TraceIn_RightLimitSwitch[192] := BenchUut15.RightLimitSwitch;
   TraceIn_GripLimitSwitch[192] := BenchUut15.GripLimitSwitch;
   TraceIn_ReleaseLimitSwitch[192] := BenchUut15.ReleaseLimitSwitch;
   BenchUut15();
   TraceOut_MoveDown[192] := BenchUut15.MoveDown;
   TraceOut_MoveUp[192] := BenchUut15.MoveUp;
   TraceOut_MoveLeft[192] := BenchUut15.MoveLeft;
   TraceOut_MoveRight[192] := BenchUut15.MoveRight;
   TraceOut_ActivateGrip[192] := BenchUut15.ActivateGrip;
   TraceOut_ActivateRelease[192] := BenchUut15.ActivateRelease;
   BenchCalls := BenchCalls + 1;
 193:
   BenchUut15.ManualMode := FALSE;
   BenchUut15.SingleStepMode := FALSE;
   BenchUut15.SingleCycleMode := TRUE;
   BenchUut15.ContinuousMode := FALSE;
   BenchUut15.EmergencyStop := TRUE;
   BenchUut15.Start := FALSE;
   BenchUut15.DownButton := FALSE;
   BenchUut15.UpButton := FALSE;
   BenchUut15.LeftButton := FALSE;
   BenchUut15.RightButton := FALSE;
   BenchUut15.GripButton := FALSE;
   BenchUut15.ReleaseButton := FALSE;
   BenchUut15.DownLimitSwitch := FALSE;
   BenchUut15.UpLimitSwitch := FALSE;
   BenchUut15.LeftLimitSwitch := FALSE;
   BenchUut15.RightLimitSwitch := FALSE;
   BenchUut15.GripLimitSwitch := FALSE;
   BenchUut15.ReleaseLimitSwitch := FALSE;
   TraceIn_ManualMode[193] := BenchUut15.ManualMode;
   TraceIn_SingleStepMode[193] := BenchUut15.SingleStepMode;
   TraceIn_SingleCycleMode[193] := BenchUut15.SingleCycleMode;
   TraceIn_ContinuousMode[193] := BenchUut15.ContinuousMode;
   TraceIn_EmergencyStop[193] := BenchUut15.EmergencyStop;
   TraceIn_Sta